(* IEC 61131-3 sources: plc-hackathon-2026/work/dump/MyController/Plc Logic/Application/Init (part 4) *)

(* ---- Init_Prof_PriceDA.st ---- *)
FUNCTION_BLOCK Init_Prof_PriceDA
VAR_INPUT
END_VAR
VAR_OUTPUT
END_VAR
VAR
END_VAR

// ---IMPL---
// Inicijalizacija GVL "Prof_PriceDA"
   Prof_PriceDA.Data[0] := 0.1353348;
   Prof_PriceDA.Data[1] := 0.1353348;
   Prof_PriceDA.Data[2] := 0.1353348;
   Prof_PriceDA.Data[3] := 0.1353348;
   Prof_PriceDA.Data[4] := 0.143694;
   Prof_PriceDA.Data[5] := 0.143694;
   Prof_PriceDA.Data[6] := 0.143694;
   Prof_PriceDA.Data[7] := 0.143694;
   Prof_PriceDA.Data[8] := 0.1349352;
   Prof_PriceDA.Data[9] := 0.1349352;
   Prof_PriceDA.Data[10] := 0.1349352;
   Prof_PriceDA.Data[11] := 0.1349352;
   Prof_PriceDA.Data[12] := 0.1010124;
   Prof_PriceDA.Data[13] := 0.1010124;
   Prof_PriceDA.Data[14] := 0.1010124;
   Prof_PriceDA.Data[15] := 0.1010124;
   Prof_PriceDA.Data[16] := 0.0687852;
   Prof_PriceDA.Data[17] := 0.0687852;
   Prof_PriceDA.Data[18] := 0.0687852;
   Prof_PriceDA.Data[19] := 0.0687852;
   Prof_PriceDA.Data[20] := 0.1011852;
   Prof_PriceDA.Data[21] := 0.1011852;
   Prof_PriceDA.Data[22] := 0.1011852;
   Prof_PriceDA.Data[23] := 0.1011852;
   Prof_PriceDA.Data[24] := 0.0974808;
   Prof_PriceDA.Data[25] := 0.0974808;
   Prof_PriceDA.Data[26] := 0.0974808;
   Prof_PriceDA.Data[27] := 0.0974808;
   Prof_PriceDA.Data[28] := 0.0902556;
   Prof_PriceDA.Data[29] := 0.0902556;
   Prof_PriceDA.Data[30] := 0.0902556;
   Prof_PriceDA.Data[31] := 0.0902556;
   Prof_PriceDA.Data[32] := 0.0399492;
   Prof_PriceDA.Data[33] := 0.0399492;
   Prof_PriceDA.Data[34] := 0.0399492;
   Prof_PriceDA.Data[35] := 0.0399492;
   Prof_PriceDA.Data[36] := 0.0485892;
   Prof_PriceDA.Data[37] := 0.0485892;
   Prof_PriceDA.Data[38] := 0.0485892;
   Prof_PriceDA.Data[39] := 0.0485892;
   Prof_PriceDA.Data[40] := 0.04158;
   Prof_PriceDA.Data[41] := 0.04158;
   Prof_PriceDA.Data[42] := 0.04158;
   Prof_PriceDA.Data[43] := 0.04158;
   Prof_PriceDA.Data[44] := 0.0430056;
   Prof_PriceDA.Data[45] := 0.0430056;
   Prof_PriceDA.Data[46] := 0.0430056;
   Prof_PriceDA.Data[47] := 0.0430056;
   Prof_PriceDA.Data[48] := 0.04347;
   Prof_PriceDA.Data[49] := 0.04347;
   Prof_PriceDA.Data[50] := 0.04347;
   Prof_PriceDA.Data[51] := 0.04347;
   Prof_PriceDA.Data[52] := 0.059886;
   Prof_PriceDA.Data[53] := 0.059886;
   Prof_PriceDA.Data[54] := 0.059886;
   Prof_PriceDA.Data[55] := 0.059886;
   Prof_PriceDA.Data[56] := 0.0664632;
   Prof_PriceDA.Data[57] := 0.0664632;
   Prof_PriceDA.Data[58] := 0.0664632;
   Prof_PriceDA.Data[59] := 0.0664632;
   Prof_PriceDA.Data[60] := 0.0900288;
   Prof_PriceDA.Data[61] := 0.0900288;
   Prof_PriceDA.Data[62] := 0.0900288;
   Prof_PriceDA.Data[63] := 0.0900288;
   Prof_PriceDA.Data[64] := 0.1161648;
   Prof_PriceDA.Data[65] := 0.1161648;
   Prof_PriceDA.Data[66] := 0.1161648;
   Prof_PriceDA.Data[67] := 0.1161648;
   Prof_PriceDA.Data[68] := 0.1328832;
   Prof_PriceDA.Data[69] := 0.1328832;
   Prof_PriceDA.Data[70] := 0.1328832;
   Prof_PriceDA.Data[71] := 0.1328832;
   Prof_PriceDA.Data[72] := 0.1382724;
   Prof_PriceDA.Data[73] := 0.1382724;
   Prof_PriceDA.Data[74] := 0.1382724;
   Prof_PriceDA.Data[75] := 0.1382724;
   Prof_PriceDA.Data[76] := 0.1446984;
   Prof_PriceDA.Data[77] := 0.1446984;
   Prof_PriceDA.Data[78] := 0.1446984;
   Prof_PriceDA.Data[79] := 0.1446984;
   Prof_PriceDA.Data[80] := 0.1406268;
   Prof_PriceDA.Data[81] := 0.1406268;
   Prof_PriceDA.Data[82] := 0.1406268;
   Prof_PriceDA.Data[83] := 0.1406268;
   Prof_PriceDA.Data[84] := 0.1307124;
   Prof_PriceDA.Data[85] := 0.1307124;
   Prof_PriceDA.Data[86] := 0.1307124;
   Prof_PriceDA.Data[87] := 0.1307124;
   Prof_PriceDA.Data[88] := 0.1310364;
   Prof_PriceDA.Data[89] := 0.1310364;
   Prof_PriceDA.Data[90] := 0.1310364;
   Prof_PriceDA.Data[91] := 0.1310364;
   Prof_PriceDA.Data[92] := 0.0904176;
   Prof_PriceDA.Data[93] := 0.0904176;
   Prof_PriceDA.Data[94] := 0.0904176;
   Prof_PriceDA.Data[95] := 0.0904176;
   Prof_PriceDA.Data[96] := 0.0689904;
   Prof_PriceDA.Data[97] := 0.0689904;
   Prof_PriceDA.Data[98] := 0.0689904;
   Prof_PriceDA.Data[99] := 0.0689904;
   Prof_PriceDA.Data[100] := 0.0865296;
   Prof_PriceDA.Data[101] := 0.0865296;
   Prof_PriceDA.Data[102] := 0.0865296;
   Prof_PriceDA.Data[103] := 0.0865296;
   Prof_PriceDA.Data[104] := 0.0846936;
   Prof_PriceDA.Data[105] := 0.0846936;
   Prof_PriceDA.Data[106] := 0.0846936;
   Prof_PriceDA.Data[107] := 0.0846936;
   Prof_PriceDA.Data[108] := 0.053136;
   Prof_PriceDA.Data[109] := 0.053136;
   Prof_PriceDA.Data[110] := 0.053136;
   Prof_PriceDA.Data[111] := 0.053136;
   Prof_PriceDA.Data[112] := 0.0614844;
   Prof_PriceDA.Data[113] := 0.0614844;
   Prof_PriceDA.Data[114] := 0.0614844;
   Prof_PriceDA.Data[115] := 0.0614844;
   Prof_PriceDA.Data[116] := 0.0834732;
   Prof_PriceDA.Data[117] := 0.0834732;
   Prof_PriceDA.Data[118] := 0.0834732;
   Prof_PriceDA.Data[119] := 0.0834732;
   Prof_PriceDA.Data[120] := 0.1200204;
   Prof_PriceDA.Data[121] := 0.1200204;
   Prof_PriceDA.Data[122] := 0.1200204;
   Prof_PriceDA.Data[123] := 0.1200204;
   Prof_PriceDA.Data[124] := 0.1431324;
   Prof_PriceDA.Data[125] := 0.1431324;
   Prof_PriceDA.Data[126] := 0.1431324;
   Prof_PriceDA.Data[127] := 0.1431324;
   Prof_PriceDA.Data[128] := 0.1405836;
   Prof_PriceDA.Data[129] := 0.1405836;
   Prof_PriceDA.Data[130] := 0.1405836;
   Prof_PriceDA.Data[131] := 0.1405836;
   Prof_PriceDA.Data[132] := 0.1433268;
   Prof_PriceDA.Data[133] := 0.1433268;
   Prof_PriceDA.Data[134] := 0.1433268;
   Prof_PriceDA.Data[135] := 0.1433268;
   Prof_PriceDA.Data[136] := 0.1391148;
   Prof_PriceDA.Data[137] := 0.1391148;
   Prof_PriceDA.Data[138] := 0.1391148;
   Prof_PriceDA.Data[139] := 0.1391148;
   Prof_PriceDA.Data[140] := 0.1337364;
   Prof_PriceDA.Data[141] := 0.1337364;
   Prof_PriceDA.Data[142] := 0.1337364;
   Prof_PriceDA.Data[143] := 0.1337364;
   Prof_PriceDA.Data[144] := 0.1330668;
   Prof_PriceDA.Data[145] := 0.1330668;
   Prof_PriceDA.Data[146] := 0.1330668;
   Prof_PriceDA.Data[147] := 0.1330668;
   Prof_PriceDA.Data[148] := 0.126144;
   Prof_PriceDA.Data[149] := 0.126144;
   Prof_PriceDA.Data[150] := 0.126144;
   Prof_PriceDA.Data[151] := 0.126144;
   Prof_PriceDA.Data[152] := 0.135;
   Prof_PriceDA.Data[153] := 0.135;
   Prof_PriceDA.Data[154] := 0.135;
   Prof_PriceDA.Data[155] := 0.135;
   Prof_PriceDA.Data[156] := 0.1405188;
   Prof_PriceDA.Data[157] := 0.1405188;
   Prof_PriceDA.Data[158] := 0.1405188;
   Prof_PriceDA.Data[159] := 0.1405188;
   Prof_PriceDA.Data[160] := 0.1650456;
   Prof_PriceDA.Data[161] := 0.1650456;
   Prof_PriceDA.Data[162] := 0.1650456;
   Prof_PriceDA.Data[163] := 0.1650456;
   Prof_PriceDA.Data[164] := 0.1762452;
   Prof_PriceDA.Data[165] := 0.1762452;
   Prof_PriceDA.Data[166] := 0.1762452;
   Prof_PriceDA.Data[167] := 0.1762452;
   Prof_PriceDA.Data[168] := 0.1695492;
   Prof_PriceDA.Data[169] := 0.1695492;
   Prof_PriceDA.Data[170] := 0.1695492;
   Prof_PriceDA.Data[171] := 0.1695492;
   Prof_PriceDA.Data[172] := 0.1646028;
   Prof_PriceDA.Data[173] := 0.1646028;
   Prof_PriceDA.Data[174] := 0.1646028;
   Prof_PriceDA.Data[175] := 0.1646028;
   Prof_PriceDA.Data[176] := 0.1414152;
   Prof_PriceDA.Data[177] := 0.1414152;
   Prof_PriceDA.Data[178] := 0.1414152;
   Prof_PriceDA.Data[179] := 0.1414152;
   Prof_PriceDA.Data[180] := 0.134622;
   Prof_PriceDA.Data[181] := 0.134622;
   Prof_PriceDA.Data[182] := 0.134622;
   Prof_PriceDA.Data[183] := 0.134622;
   Prof_PriceDA.Data[184] := 0.1270188;
   Prof_PriceDA.Data[185] := 0.1270188;
   Prof_PriceDA.Data[186] := 0.1270188;
   Prof_PriceDA.Data[187] := 0.1270188;
   Prof_PriceDA.Data[188] := 0.1095228;
   Prof_PriceDA.Data[189] := 0.1095228;
   Prof_PriceDA.Data[190] := 0.1095228;
   Prof_PriceDA.Data[191] := 0.1095228;
   Prof_PriceDA.Data[192] := 0.111996;
   Prof_PriceDA.Data[193] := 0.111996;
   Prof_PriceDA.Data[194] := 0.111996;
   Prof_PriceDA.Data[195] := 0.111996;
   Prof_PriceDA.Data[196] := 0.1023732;
   Prof_PriceDA.Data[197] := 0.1023732;
   Prof_PriceDA.Data[198] := 0.1023732;
   Prof_PriceDA.Data[199] := 0.1023732;
   Prof_PriceDA.Data[200] := 0.0968436;
   Prof_PriceDA.Data[201] := 0.0968436;
   Prof_PriceDA.Data[202] := 0.0968436;
   Prof_PriceDA.Data[203] := 0.0968436;
   Prof_PriceDA.Data[204] := 0.0945216;
   Prof_PriceDA.Data[205] := 0.0945216;
   Prof_PriceDA.Data[206] := 0.0945216;
   Prof_PriceDA.Data[207] := 0.0945216;
   Prof_PriceDA.Data[208] := 0.0923832;
   Prof_PriceDA.Data[209] := 0.0923832;
   Prof_PriceDA.Data[210] := 0.0923832;
   Prof_PriceDA.Data[211] := 0.0923832;
   Prof_PriceDA.Data[212] := 0.0993816;
   Prof_PriceDA.Data[213] := 0.0993816;
   Prof_PriceDA.Data[214] := 0.0993816;
   Prof_PriceDA.Data[215] := 0.0993816;
   Prof_PriceDA.Data[216] := 0.1185516;
   Prof_PriceDA.Data[217] := 0.1185516;
   Prof_PriceDA.Data[218] := 0.1185516;
   Prof_PriceDA.Data[219] := 0.1185516;
   Prof_PriceDA.Data[220] := 0.1469556;
   Prof_PriceDA.Data[221] := 0.1469556;
   Prof_PriceDA.Data[222] := 0.1469556;
   Prof_PriceDA.Data[223] := 0.1469556;
   Prof_PriceDA.Data[224] := 0.1492452;
   Prof_PriceDA.Data[225] := 0.1492452;
   Prof_PriceDA.Data[226] := 0.1492452;
   Prof_PriceDA.Data[227] := 0.1492452;
   Prof_PriceDA.Data[228] := 0.1461564;
   Prof_PriceDA.Data[229] := 0.1461564;
   Prof_PriceDA.Data[230] := 0.1461564;
   Prof_PriceDA.Data[231] := 0.1461564;
   Prof_PriceDA.Data[232] := 0.1350216;
   Prof_PriceDA.Data[233] := 0.1350216;
   Prof_PriceDA.Data[234] := 0.1350216;
   Prof_PriceDA.Data[235] := 0.1350216;
   Prof_PriceDA.Data[236] := 0.1219968;
   Prof_PriceDA.Data[237] := 0.1219968;
   Prof_PriceDA.Data[238] := 0.1219968;
   Prof_PriceDA.Data[239] := 0.1219968;
   Prof_PriceDA.Data[240] := 0.1201716;
   Prof_PriceDA.Data[241] := 0.1201716;
   Prof_PriceDA.Data[242] := 0.1201716;
   Prof_PriceDA.Data[243] := 0.1201716;
   Prof_PriceDA.Data[244] := 0.118206;
   Prof_PriceDA.Data[245] := 0.118206;
   Prof_PriceDA.Data[246] := 0.118206;
   Prof_PriceDA.Data[247] := 0.118206;
   Prof_PriceDA.Data[248] := 0.124956;
   Prof_PriceDA.Data[249] := 0.124956;
   Prof_PriceDA.Data[250] := 0.124956;
   Prof_PriceDA.Data[251] := 0.124956;
   Prof_PriceDA.Data[252] := 0.1402596;
   Prof_PriceDA.Data[253] := 0.1402596;
   Prof_PriceDA.Data[254] := 0.1402596;
   Prof_PriceDA.Data[255] := 0.1402596;
   Prof_PriceDA.Data[256] := 0.1587276;
   Prof_PriceDA.Data[257] := 0.1587276;
   Prof_PriceDA.Data[258] := 0.1587276;
   Prof_PriceDA.Data[259] := 0.1587276;
   Prof_PriceDA.Data[260] := 0.1571508;
   Prof_PriceDA.Data[261] := 0.1571508;
   Prof_PriceDA.Data[262] := 0.1571508;
   Prof_PriceDA.Data[263] := 0.1571508;
   Prof_PriceDA.Data[264] := 0.1572696;
   Prof_PriceDA.Data[265] := 0.1572696;
   Prof_PriceDA.Data[266] := 0.1572696;
   Prof_PriceDA.Data[267] := 0.1572696;
   Prof_PriceDA.Data[268] := 0.1564488;
   Prof_PriceDA.Data[269] := 0.1564488;
   Prof_PriceDA.Data[270] := 0.1564488;
   Prof_PriceDA.Data[271] := 0.1564488;
   Prof_PriceDA.Data[272] := 0.1478196;
   Prof_PriceDA.Data[273] := 0.1478196;
   Prof_PriceDA.Data[274] := 0.1478196;
   Prof_PriceDA.Data[275] := 0.1478196;
   Prof_PriceDA.Data[276] := 0.1314684;
   Prof_PriceDA.Data[277] := 0.1314684;
   Prof_PriceDA.Data[278] := 0.1314684;
   Prof_PriceDA.Data[279] := 0.1314684;
   Prof_PriceDA.Data[280] := 0.1361988;
   Prof_PriceDA.Data[281] := 0.1361988;
   Prof_PriceDA.Data[282] := 0.1361988;
   Prof_PriceDA.Data[283] := 0.1361988;
   Prof_PriceDA.Data[284] := 0.1318572;
   Prof_PriceDA.Data[285] := 0.1318572;
   Prof_PriceDA.Data[286] := 0.1318572;
   Prof_PriceDA.Data[287] := 0.1318572;
   Prof_PriceDA.Data[288] := 0.1189296;
   Prof_PriceDA.Data[289] := 0.1189296;
   Prof_PriceDA.Data[290] := 0.1189296;
   Prof_PriceDA.Data[291] := 0.1189296;
   Prof_PriceDA.Data[292] := 0.1130112;
   Prof_PriceDA.Data[293] := 0.1130112;
   Prof_PriceDA.Data[294] := 0.1130112;
   Prof_PriceDA.Data[295] := 0.1130112;
   Prof_PriceDA.Data[296] := 0.1087344;
   Prof_PriceDA.Data[297] := 0.1087344;
   Prof_PriceDA.Data[298] := 0.1087344;
   Prof_PriceDA.Data[299] := 0.1087344;
   Prof_PriceDA.Data[300] := 0.1065204;
   Prof_PriceDA.Data[301] := 0.1065204;
   Prof_PriceDA.Data[302] := 0.1065204;
   Prof_PriceDA.Data[303] := 0.1065204;
   Prof_PriceDA.Data[304] := 0.1077732;
   Prof_PriceDA.Data[305] := 0.1077732;
   Prof_PriceDA.Data[306] := 0.1077732;
   Prof_PriceDA.Data[307] := 0.1077732;
   Prof_PriceDA.Data[308] := 0.113454;
   Prof_PriceDA.Data[309] := 0.113454;
   Prof_PriceDA.Data[310] := 0.113454;
   Prof_PriceDA.Data[311] := 0.113454;
   Prof_PriceDA.Data[312] := 0.12096;
   Prof_PriceDA.Data[313] := 0.12096;
   Prof_PriceDA.Data[314] := 0.12096;
   Prof_PriceDA.Data[315] := 0.12096;
   Prof_PriceDA.Data[316] := 0.1352808;
   Prof_PriceDA.Data[317] := 0.1352808;
   Prof_PriceDA.Data[318] := 0.1352808;
   Prof_PriceDA.Data[319] := 0.1352808;
   Prof_PriceDA.Data[320] := 0.1386612;
   Prof_PriceDA.Data[321] := 0.1386612;
   Prof_PriceDA.Data[322] := 0.1386612;
   Prof_PriceDA.Data[323] := 0.1386612;
   Prof_PriceDA.Data[324] := 0.14121;
   Prof_PriceDA.Data[325] := 0.14121;
   Prof_PriceDA.Data[326] := 0.14121;
   Prof_PriceDA.Data[327] := 0.14121;
   Prof_PriceDA.Data[328] := 0.1407672;
   Prof_PriceDA.Data[329] := 0.1407672;
   Prof_PriceDA.Data[330] := 0.1407672;
   Prof_PriceDA.Data[331] := 0.1407672;
   Prof_PriceDA.Data[332] := 0.1385532;
   Prof_PriceDA.Data[333] := 0.1385532;
   Prof_PriceDA.Data[334] := 0.1385532;
   Prof_PriceDA.Data[335] := 0.1385532;
   Prof_PriceDA.Data[336] := 0.1404324;
   Prof_PriceDA.Data[337] := 0.1404324;
   Prof_PriceDA.Data[338] := 0.1404324;
   Prof_PriceDA.Data[339] := 0.1404324;
   Prof_PriceDA.Data[340] := 0.140238;
   Prof_PriceDA.Data[341] := 0.140238;
   Prof_PriceDA.Data[342] := 0.140238;
   Prof_PriceDA.Data[343] := 0.140238;
   Prof_PriceDA.Data[344] := 0.147312;
   Prof_PriceDA.Data[345] := 0.147312;
   Prof_PriceDA.Data[346] := 0.147312;
   Prof_PriceDA.Data[347] := 0.147312;
   Prof_PriceDA.Data[348] := 0.15309;
   Prof_PriceDA.Data[349] := 0.15309;
   Prof_PriceDA.Data[350] := 0.15309;
   Prof_PriceDA.Data[351] := 0.15309;
   Prof_PriceDA.Data[352] := 0.1819368;
   Prof_PriceDA.Data[353] := 0.1819368;
   Prof_PriceDA.Data[354] := 0.1819368;
   Prof_PriceDA.Data[355] := 0.1819368;
   Prof_PriceDA.Data[356] := 0.1857924;
   Prof_PriceDA.Data[357] := 0.1857924;
   Prof_PriceDA.Data[358] := 0.1857924;
   Prof_PriceDA.Data[359] := 0.1857924;
   Prof_PriceDA.Data[360] := 0.1848096;
   Prof_PriceDA.Data[361] := 0.1848096;
   Prof_PriceDA.Data[362] := 0.1848096;
   Prof_PriceDA.Data[363] := 0.1848096;
   Prof_PriceDA.Data[364] := 0.1831572;
   Prof_PriceDA.Data[365] := 0.1831572;
   Prof_PriceDA.Data[366] := 0.1831572;
   Prof_PriceDA.Data[367] := 0.1831572;
   Prof_PriceDA.Data[368] := 0.1590624;
   Prof_PriceDA.Data[369] := 0.1590624;
   Prof_PriceDA.Data[370] := 0.1590624;
   Prof_PriceDA.Data[371] := 0.1590624;
   Prof_PriceDA.Data[372] := 0.151524;
   Prof_PriceDA.Data[373] := 0.151524;
   Prof_PriceDA.Data[374] := 0.151524;
   Prof_PriceDA.Data[375] := 0.151524;
   Prof_PriceDA.Data[376] := 0.1455192;
   Prof_PriceDA.Data[377] := 0.1455192;
   Prof_PriceDA.Data[378] := 0.1455192;
   Prof_PriceDA.Data[379] := 0.1455192;
   Prof_PriceDA.Data[380] := 0.1259604;
   Prof_PriceDA.Data[381] := 0.1259604;
   Prof_PriceDA.Data[382] := 0.1259604;
   Prof_PriceDA.Data[383] := 0.1259604;
   Prof_PriceDA.Data[384] := 0.1211004;
   Prof_PriceDA.Data[385] := 0.1211004;
   Prof_PriceDA.Data[386] := 0.1211004;
   Prof_PriceDA.Data[387] := 0.1211004;
   Prof_PriceDA.Data[388] := 0.107838;
   Prof_PriceDA.Data[389] := 0.107838;
   Prof_PriceDA.Data[390] := 0.107838;
   Prof_PriceDA.Data[391] := 0.107838;
   Prof_PriceDA.Data[392] := 0.1033668;
   Prof_PriceDA.Data[393] := 0.1033668;
   Prof_PriceDA.Data[394] := 0.1033668;
   Prof_PriceDA.Data[395] := 0.1033668;
   Prof_PriceDA.Data[396] := 0.1013364;
   Prof_PriceDA.Data[397] := 0.1013364;
   Prof_PriceDA.Data[398] := 0.1013364;
   Prof_PriceDA.Data[399] := 0.1013364;
   Prof_PriceDA.Data[400] := 0.1006992;
   Prof_PriceDA.Data[401] := 0.1006992;
   Prof_PriceDA.Data[402] := 0.1006992;
   Prof_PriceDA.Data[403] := 0.1006992;
   Prof_PriceDA.Data[404] := 0.0971892;
   Prof_PriceDA.Data[405] := 0.0971892;
   Prof_PriceDA.Data[406] := 0.0971892;
   Prof_PriceDA.Data[407] := 0.0971892;
   Prof_PriceDA.Data[408] := 0.0989064;
   Prof_PriceDA.Data[409] := 0.0989064;
   Prof_PriceDA.Data[410] := 0.0989064;
   Prof_PriceDA.Data[411] := 0.0989064;
   Prof_PriceDA.Data[412] := 0.1068012;
   Prof_PriceDA.Data[413] := 0.1068012;
   Prof_PriceDA.Data[414] := 0.1068012;
   Prof_PriceDA.Data[415] := 0.1068012;
   Prof_PriceDA.Data[416] := 0.105408;
   Prof_PriceDA.Data[417] := 0.105408;
   Prof_PriceDA.Data[418] := 0.105408;
   Prof_PriceDA.Data[419] := 0.105408;
   Prof_PriceDA.Data[420] := 0.1070172;
   Prof_PriceDA.Data[421] := 0.1070172;
   Prof_PriceDA.Data[422] := 0.1070172;
   Prof_PriceDA.Data[423] := 0.1070172;
   Prof_PriceDA.Data[424] := 0.103194;
   Prof_PriceDA.Data[425] := 0.103194;
   Prof_PriceDA.Data[426] := 0.103194;
   Prof_PriceDA.Data[427] := 0.103194;
   Prof_PriceDA.Data[428] := 0.1084104;
   Prof_PriceDA.Data[429] := 0.1084104;
   Prof_PriceDA.Data[430] := 0.1084104;
   Prof_PriceDA.Data[431] := 0.1084104;
   Prof_PriceDA.Data[432] := 0.1057752;
   Prof_PriceDA.Data[433] := 0.1057752;
   Prof_PriceDA.Data[434] := 0.1057752;
   Prof_PriceDA.Data[435] := 0.1057752;
   Prof_PriceDA.Data[436] := 0.1129248;
   Prof_PriceDA.Data[437] := 0.1129248;
   Prof_PriceDA.Data[438] := 0.1129248;
   Prof_PriceDA.Data[439] := 0.1129248;
   Prof_PriceDA.Data[440] := 0.122094;
   Prof_PriceDA.Data[441] := 0.122094;
   Prof_PriceDA.Data[442] := 0.122094;
   Prof_PriceDA.Data[443] := 0.122094;
   Prof_PriceDA.Data[444] := 0.1337364;
   Prof_PriceDA.Data[445] := 0.1337364;
   Prof_PriceDA.Data[446] := 0.1337364;
   Prof_PriceDA.Data[447] := 0.1337364;
   Prof_PriceDA.Data[448] := 0.1717308;
   Prof_PriceDA.Data[449] := 0.1717308;
   Prof_PriceDA.Data[450] := 0.1717308;
   Prof_PriceDA.Data[451] := 0.1717308;
   Prof_PriceDA.Data[452] := 0.165024;
   Prof_PriceDA.Data[453] := 0.165024;
   Prof_PriceDA.Data[454] := 0.165024;
   Prof_PriceDA.Data[455] := 0.165024;
   Prof_PriceDA.Data[456] := 0.1562328;
   Prof_PriceDA.Data[457] := 0.1562328;
   Prof_PriceDA.Data[458] := 0.1562328;
   Prof_PriceDA.Data[459] := 0.1562328;
   Prof_PriceDA.Data[460] := 0.1627236;
   Prof_PriceDA.Data[461] := 0.1627236;
   Prof_PriceDA.Data[462] := 0.1627236;
   Prof_PriceDA.Data[463] := 0.1627236;
   Prof_PriceDA.Data[464] := 0.1535328;
   Prof_PriceDA.Data[465] := 0.1535328;
   Prof_PriceDA.Data[466] := 0.1535328;
   Prof_PriceDA.Data[467] := 0.1535328;
   Prof_PriceDA.Data[468] := 0.1449144;
   Prof_PriceDA.Data[469] := 0.1449144;
   Prof_PriceDA.Data[470] := 0.1449144;
   Prof_PriceDA.Data[471] := 0.1449144;
   Prof_PriceDA.Data[472] := 0.1105056;
   Prof_PriceDA.Data[473] := 0.1105056;
   Prof_PriceDA.Data[474] := 0.1105056;
   Prof_PriceDA.Data[475] := 0.1105056;
   Prof_PriceDA.Data[476] := 0.0771984;
   Prof_PriceDA.Data[477] := 0.0771984;
   Prof_PriceDA.Data[478] := 0.0771984;
   Prof_PriceDA.Data[479] := 0.0771984;
   Prof_PriceDA.Data[480] := 0.1130004;
   Prof_PriceDA.Data[481] := 0.1130004;
   Prof_PriceDA.Data[482] := 0.1130004;
   Prof_PriceDA.Data[483] := 0.1130004;
   Prof_PriceDA.Data[484] := 0.0960336;
   Prof_PriceDA.Data[485] := 0.0960336;
   Prof_PriceDA.Data[486] := 0.0960336;
   Prof_PriceDA.Data[487] := 0.0960336;
   Prof_PriceDA.Data[488] := 0.0743256;
   Prof_PriceDA.Data[489] := 0.0743256;
   Prof_PriceDA.Data[490] := 0.0743256;
   Prof_PriceDA.Data[491] := 0.0743256;
   Prof_PriceDA.Data[492] := 0.0708804;
   Prof_PriceDA.Data[493] := 0.0708804;
   Prof_PriceDA.Data[494] := 0.0708804;
   Prof_PriceDA.Data[495] := 0.0708804;
   Prof_PriceDA.Data[496] := 0.070794;
   Prof_PriceDA.Data[497] := 0.070794;
   Prof_PriceDA.Data[498] := 0.070794;
   Prof_PriceDA.Data[499] := 0.070794;
   Prof_PriceDA.Data[500] := 0.0962172;
   Prof_PriceDA.Data[501] := 0.0962172;
   Prof_PriceDA.Data[502] := 0.0962172;
   Prof_PriceDA.Data[503] := 0.0962172;
   Prof_PriceDA.Data[504] := 0.1229364;
   Prof_PriceDA.Data[505] := 0.1229364;
   Prof_PriceDA.Data[506] := 0.1229364;
   Prof_PriceDA.Data[507] := 0.1229364;
   Prof_PriceDA.Data[508] := 0.1331748;
   Prof_PriceDA.Data[509] := 0.1331748;
   Prof_PriceDA.Data[510] := 0.1331748;
   Prof_PriceDA.Data[511] := 0.1331748;
   Prof_PriceDA.Data[512] := 0.1334664;
   Prof_PriceDA.Data[513] := 0.1334664;
   Prof_PriceDA.Data[514] := 0.1334664;
   Prof_PriceDA.Data[515] := 0.1334664;
   Prof_PriceDA.Data[516] := 0.1152576;
   Prof_PriceDA.Data[517] := 0.1152576;
   Prof_PriceDA.Data[518] := 0.1152576;
   Prof_PriceDA.Data[519] := 0.1152576;
   Prof_PriceDA.Data[520] := 0.097956;
   Prof_PriceDA.Data[521] := 0.097956;
   Prof_PriceDA.Data[522] := 0.097956;
   Prof_PriceDA.Data[523] := 0.097956;
   Prof_PriceDA.Data[524] := 0.0780624;
   Prof_PriceDA.Data[525] := 0.0780624;
   Prof_PriceDA.Data[526] := 0.0780624;
   Prof_PriceDA.Data[527] := 0.0780624;
   Prof_PriceDA.Data[528] := 0.0841212;
   Prof_PriceDA.Data[529] := 0.0841212;
   Prof_PriceDA.Data[530] := 0.0841212;
   Prof_PriceDA.Data[531] := 0.0841212;
   Prof_PriceDA.Data[532] := 0.10476;
   Prof_PriceDA.Data[533] := 0.10476;
   Prof_PriceDA.Data[534] := 0.10476;
   Prof_PriceDA.Data[535] := 0.10476;
   Prof_PriceDA.Data[536] := 0.1249668;
   Prof_PriceDA.Data[537] := 0.1249668;
   Prof_PriceDA.Data[538] := 0.1249668;
   Prof_PriceDA.Data[539] := 0.1249668;
   Prof_PriceDA.Data[540] := 0.1229904;
   Prof_PriceDA.Data[541] := 0.1229904;
   Prof_PriceDA.Data[542] := 0.1229904;
   Prof_PriceDA.Data[543] := 0.1229904;
   Prof_PriceDA.Data[544] := 0.1472904;
   Prof_PriceDA.Data[545] := 0.1472904;
   Prof_PriceDA.Data[546] := 0.1472904;
   Prof_PriceDA.Data[547] := 0.1472904;
   Prof_PriceDA.Data[548] := 0.1600344;
   Prof_PriceDA.Data[549] := 0.1600344;
   Prof_PriceDA.Data[550] := 0.1600344;
   Prof_PriceDA.Data[551] := 0.1600344;
   Prof_PriceDA.Data[552] := 0.1528524;
   Prof_PriceDA.Data[553] := 0.1528524;
   Prof_PriceDA.Data[554] := 0.1528524;
   Prof_PriceDA.Data[555] := 0.1528524;
   Prof_PriceDA.Data[556] := 0.1521828;
   Prof_PriceDA.Data[557] := 0.1521828;
   Prof_PriceDA.Data[558] := 0.1521828;
   Prof_PriceDA.Data[559] := 0.1521828;
   Prof_PriceDA.Data[560] := 0.1456272;
   Prof_PriceDA.Data[561] := 0.1456272;
   Prof_PriceDA.Data[562] := 0.1456272;
   Prof_PriceDA.Data[563] := 0.1456272;
   Prof_PriceDA.Data[564] := 0.122364;
   Prof_PriceDA.Data[565] := 0.122364;
   Prof_PriceDA.Data[566] := 0.122364;
   Prof_PriceDA.Data[567] := 0.122364;
   Prof_PriceDA.Data[568] := 0.1168128;
   Prof_PriceDA.Data[569] := 0.1168128;
   Prof_PriceDA.Data[570] := 0.1168128;
   Prof_PriceDA.Data[571] := 0.1168128;
   Prof_PriceDA.Data[572] := 0.0853416;
   Prof_PriceDA.Data[573] := 0.0853416;
   Prof_PriceDA.Data[574] := 0.0853416;
   Prof_PriceDA.Data[575] := 0.0853416;
   Prof_PriceDA.Data[576] := 0.0343116;
   Prof_PriceDA.Data[577] := 0.0343116;
   Prof_PriceDA.Data[578] := 0.0343116;
   Prof_PriceDA.Data[579] := 0.0343116;
   Prof_PriceDA.Data[580] := 0.056538;
   Prof_PriceDA.Data[581] := 0.056538;
   Prof_PriceDA.Data[582] := 0.056538;
   Prof_PriceDA.Data[583] := 0.056538;
   Prof_PriceDA.Data[584] := 0.0510192;
   Prof_PriceDA.Data[585] := 0.0510192;
   Prof_PriceDA.Data[586] := 0.0510192;
   Prof_PriceDA.Data[587] := 0.0510192;
   Prof_PriceDA.Data[588] := 0.0135;
   Prof_PriceDA.Data[589] := 0.0135;
   Prof_PriceDA.Data[590] := 0.0135;
   Prof_PriceDA.Data[591] := 0.0135;
   Prof_PriceDA.Data[592] := 0.0662688;
   Prof_PriceDA.Data[593] := 0.0662688;
   Prof_PriceDA.Data[594] := 0.0662688;
   Prof_PriceDA.Data[595] := 0.0662688;
   Prof_PriceDA.Data[596] := 0.0844668;
   Prof_PriceDA.Data[597] := 0.0844668;
   Prof_PriceDA.Data[598] := 0.0844668;
   Prof_PriceDA.Data[599] := 0.0844668;
   Prof_PriceDA.Data[600] := 0.1362636;
   Prof_PriceDA.Data[601] := 0.1362636;
   Prof_PriceDA.Data[602] := 0.1362636;
   Prof_PriceDA.Data[603] := 0.1362636;
   Prof_PriceDA.Data[604] := 0.16443;
   Prof_PriceDA.Data[605] := 0.16443;
   Prof_PriceDA.Data[606] := 0.16443;
   Prof_PriceDA.Data[607] := 0.16443;
   Prof_PriceDA.Data[608] := 0.148014;
   Prof_PriceDA.Data[609] := 0.148014;
   Prof_PriceDA.Data[610] := 0.148014;
   Prof_PriceDA.Data[611] := 0.148014;
   Prof_PriceDA.Data[612] := 0.1423224;
   Prof_PriceDA.Data[613] := 0.1423224;
   Prof_PriceDA.Data[614] := 0.1423224;
   Prof_PriceDA.Data[615] := 0.1423224;
   Prof_PriceDA.Data[616] := 0.1318248;
   Prof_PriceDA.Data[617] := 0.1318248;
   Prof_PriceDA.Data[618] := 0.1318248;
   Prof_PriceDA.Data[619] := 0.1318248;
   Prof_PriceDA.Data[620] := 0.131274;
   Prof_PriceDA.Data[621] := 0.131274;
   Prof_PriceDA.Data[622] := 0.131274;
   Prof_PriceDA.Data[623] := 0.131274;
   Prof_PriceDA.Data[624] := 0.1322676;
   Prof_PriceDA.Data[625] := 0.1322676;
   Prof_PriceDA.Data[626] := 0.1322676;
   Prof_PriceDA.Data[627] := 0.1322676;
   Prof_PriceDA.Data[628] := 0.1404432;
   Prof_PriceDA.Data[629] := 0.1404432;
   Prof_PriceDA.Data[630] := 0.1404432;
   Prof_PriceDA.Data[631] := 0.1404432;
   Prof_PriceDA.Data[632] := 0.1504656;
   Prof_PriceDA.Data[633] := 0.1504656;
   Prof_PriceDA.Data[634] := 0.1504656;
   Prof_PriceDA.Data[635] := 0.1504656;
   Prof_PriceDA.Data[636] := 0.1588572;
   Prof_PriceDA.Data[637] := 0.1588572;
   Prof_PriceDA.Data[638] := 0.1588572;
   Prof_PriceDA.Data[639] := 0.1588572;
   Prof_PriceDA.Data[640] := 0.1668384;
   Prof_PriceDA.Data[641] := 0.1668384;
   Prof_PriceDA.Data[642] := 0.1668384;
   Prof_PriceDA.Data[643] := 0.1668384;
   Prof_PriceDA.Data[644] := 0.166806;
   Prof_PriceDA.Data[645] := 0.166806;
   Prof_PriceDA.Data[646] := 0.166806;
   Prof_PriceDA.Data[647] := 0.166806;
   Prof_PriceDA.Data[648] := 0.1628424;
   Prof_PriceDA.Data[649] := 0.1628424;
   Prof_PriceDA.Data[650] := 0.1628424;
   Prof_PriceDA.Data[651] := 0.1628424;
   Prof_PriceDA.Data[652] := 0.1643328;
   Prof_PriceDA.Data[653] := 0.1643328;
   Prof_PriceDA.Data[654] := 0.1643328;
   Prof_PriceDA.Data[655] := 0.1643328;
   Prof_PriceDA.Data[656] := 0.1532088;
   Prof_PriceDA.Data[657] := 0.1532088;
   Prof_PriceDA.Data[658] := 0.1532088;
   Prof_PriceDA.Data[659] := 0.1532088;
   Prof_PriceDA.Data[660] := 0.1370196;
   Prof_PriceDA.Data[661] := 0.1370196;
   Prof_PriceDA.Data[662] := 0.1370196;
   Prof_PriceDA.Data[663] := 0.1370196;
   Prof_PriceDA.Data[664] := 0.125064;
   Prof_PriceDA.Data[665] := 0.125064;
   Prof_PriceDA.Data[666] := 0.125064;
   Prof_PriceDA.Data[667] := 0.125064;
   Prof_PriceDA.Data[668] := 0.1204416;
   Prof_PriceDA.Data[669] := 0.1204416;
   Prof_PriceDA.Data[670] := 0.1204416;
   Prof_PriceDA.Data[671] := 0.1204416;
   Prof_PriceDA.Data[672] := 0.0901584;
   Prof_PriceDA.Data[673] := 0.0901584;
   Prof_PriceDA.Data[674] := 0.0901584;
   Prof_PriceDA.Data[675] := 0.0901584;
   Prof_PriceDA.Data[676] := 0.0813672;
   Prof_PriceDA.Data[677] := 0.0813672;
   Prof_PriceDA.Data[678] := 0.0813672;
   Prof_PriceDA.Data[679] := 0.0813672;
   Prof_PriceDA.Data[680] := 0.0789048;
   Prof_PriceDA.Data[681] := 0.0789048;
   Prof_PriceDA.Data[682] := 0.0789048;
   Prof_PriceDA.Data[683] := 0.0789048;
   Prof_PriceDA.Data[684] := 0.0747036;
   Prof_PriceDA.Data[685] := 0.0747036;
   Prof_PriceDA.Data[686] := 0.0747036;
   Prof_PriceDA.Data[687] := 0.0747036;
   Prof_PriceDA.Data[688] := 0.0923076;
   Prof_PriceDA.Data[689] := 0.0923076;
   Prof_PriceDA.Data[690] := 0.0923076;
   Prof_PriceDA.Data[691] := 0.0923076;
   Prof_PriceDA.Data[692] := 0.11178;
   Prof_PriceDA.Data[693] := 0.11178;
   Prof_PriceDA.Data[694] := 0.11178;
   Prof_PriceDA.Data[695] := 0.11178;
   Prof_PriceDA.Data[696] := 0.1367388;
   Prof_PriceDA.Data[697] := 0.1367388;
   Prof_PriceDA.Data[698] := 0.1367388;
   Prof_PriceDA.Data[699] := 0.1367388;
   Prof_PriceDA.Data[700] := 0.1635336;
   Prof_PriceDA.Data[701] := 0.1635336;
   Prof_PriceDA.Data[702] := 0.1635336;
   Prof_PriceDA.Data[703] := 0.1635336;
   Prof_PriceDA.Data[704] := 0.1611252;
   Prof_PriceDA.Data[705] := 0.1611252;
   Prof_PriceDA.Data[706] := 0.1611252;
   Prof_PriceDA.Data[707] := 0.1611252;
   Prof_PriceDA.Data[708] := 0.1341576;
   Prof_PriceDA.Data[709] := 0.1341576;
   Prof_PriceDA.Data[710] := 0.1341576;
   Prof_PriceDA.Data[711] := 0.1341576;
   Prof_PriceDA.Data[712] := 0.1174068;
   Prof_PriceDA.Data[713] := 0.1174068;
   Prof_PriceDA.Data[714] := 0.1174068;
   Prof_PriceDA.Data[715] := 0.1174068;
   Prof_PriceDA.Data[716] := 0.1103436;
   Prof_PriceDA.Data[717] := 0.1103436;
   Prof_PriceDA.Data[718] := 0.1103436;
   Prof_PriceDA.Data[719] := 0.1103436;
   Prof_PriceDA.Data[720] := 0.1120824;
   Prof_PriceDA.Data[721] := 0.1120824;
   Prof_PriceDA.Data[722] := 0.1120824;
   Prof_PriceDA.Data[723] := 0.1120824;
   Prof_PriceDA.Data[724] := 0.1245996;
   Prof_PriceDA.Data[725] := 0.1245996;
   Prof_PriceDA.Data[726] := 0.1245996;
   Prof_PriceDA.Data[727] := 0.1245996;
   Prof_PriceDA.Data[728] := 0.1353132;
   Prof_PriceDA.Data[729] := 0.1353132;
   Prof_PriceDA.Data[730] := 0.1353132;
   Prof_PriceDA.Data[731] := 0.1353132;
   Prof_PriceDA.Data[732] := 0.1550556;
   Prof_PriceDA.Data[733] := 0.1550556;
   Prof_PriceDA.Data[734] := 0.1550556;
   Prof_PriceDA.Data[735] := 0.1550556;
   Prof_PriceDA.Data[736] := 0.1646784;
   Prof_PriceDA.Data[737] := 0.1646784;
   Prof_PriceDA.Data[738] := 0.1646784;
   Prof_PriceDA.Data[739] := 0.1646784;
   Prof_PriceDA.Data[740] := 0.165456;
   Prof_PriceDA.Data[741] := 0.165456;
   Prof_PriceDA.Data[742] := 0.165456;
   Prof_PriceDA.Data[743] := 0.165456;
   Prof_PriceDA.Data[744] := 0.1622916;
   Prof_PriceDA.Data[745] := 0.1622916;
   Prof_PriceDA.Data[746] := 0.1622916;
   Prof_PriceDA.Data[747] := 0.1622916;
   Prof_PriceDA.Data[748] := 0.1614384;
   Prof_PriceDA.Data[749] := 0.1614384;
   Prof_PriceDA.Data[750] := 0.1614384;
   Prof_PriceDA.Data[751] := 0.1614384;
   Prof_PriceDA.Data[752] := 0.1484352;
   Prof_PriceDA.Data[753] := 0.1484352;
   Prof_PriceDA.Data[754] := 0.1484352;
   Prof_PriceDA.Data[755] := 0.1484352;
   Prof_PriceDA.Data[756] := 0.1356372;
   Prof_PriceDA.Data[757] := 0.1356372;
   Prof_PriceDA.Data[758] := 0.1356372;
   Prof_PriceDA.Data[759] := 0.1356372;
   Prof_PriceDA.Data[760] := 0.1255716;
   Prof_PriceDA.Data[761] := 0.1255716;
   Prof_PriceDA.Data[762] := 0.1255716;
   Prof_PriceDA.Data[763] := 0.1255716;
   Prof_PriceDA.Data[764] := 0.114588;
   Prof_PriceDA.Data[765] := 0.114588;
   Prof_PriceDA.Data[766] := 0.114588;
   Prof_PriceDA.Data[767] := 0.114588;
   Prof_PriceDA.Data[768] := 0.1147284;
   Prof_PriceDA.Data[769] := 0.1147284;
   Prof_PriceDA.Data[770] := 0.1147284;
   Prof_PriceDA.Data[771] := 0.1147284;
   Prof_PriceDA.Data[772] := 0.114588;
   Prof_PriceDA.Data[773] := 0.114588;
   Prof_PriceDA.Data[774] := 0.114588;
   Prof_PriceDA.Data[775] := 0.114588;
   Prof_PriceDA.Data[776] := 0.1119096;
   Prof_PriceDA.Data[777] := 0.1119096;
   Prof_PriceDA.Data[778] := 0.1119096;
   Prof_PriceDA.Data[779] := 0.1119096;
   Prof_PriceDA.Data[780] := 0.1104408;
   Prof_PriceDA.Data[781] := 0.1104408;
   Prof_PriceDA.Data[782] := 0.1104408;
   Prof_PriceDA.Data[783] := 0.1104408;
   Prof_PriceDA.Data[784] := 0.1152468;
   Prof_PriceDA.Data[785] := 0.1152468;
   Prof_PriceDA.Data[786] := 0.1152468;
   Prof_PriceDA.Data[787] := 0.1152468;
   Prof_PriceDA.Data[788] := 0.1184868;
   Prof_PriceDA.Data[789] := 0.1184868;
   Prof_PriceDA.Data[790] := 0.1184868;
   Prof_PriceDA.Data[791] := 0.1184868;
   Prof_PriceDA.Data[792] := 0.1342656;
   Prof_PriceDA.Data[793] := 0.1342656;
   Prof_PriceDA.Data[794] := 0.1342656;
   Prof_PriceDA.Data[795] := 0.1342656;
   Prof_PriceDA.Data[796] := 0.1542132;
   Prof_PriceDA.Data[797] := 0.1542132;
   Prof_PriceDA.Data[798] := 0.1542132;
   Prof_PriceDA.Data[799] := 0.1542132;
   Prof_PriceDA.Data[800] := 0.1678104;
   Prof_PriceDA.Data[801] := 0.1678104;
   Prof_PriceDA.Data[802] := 0.1678104;
   Prof_PriceDA.Data[803] := 0.1678104;
   Prof_PriceDA.Data[804] := 0.1601208;
   Prof_PriceDA.Data[805] := 0.1601208;
   Prof_PriceDA.Data[806] := 0.1601208;
   Prof_PriceDA.Data[807] := 0.1601208;
   Prof_PriceDA.Data[808] := 0.1514916;
   Prof_PriceDA.Data[809] := 0.1514916;
   Prof_PriceDA.Data[810] := 0.1514916;
   Prof_PriceDA.Data[811] := 0.1514916;
   Prof_PriceDA.Data[812] := 0.1435644;
   Prof_PriceDA.Data[813] := 0.1435644;
   Prof_PriceDA.Data[814] := 0.1435644;
   Prof_PriceDA.Data[815] := 0.1435644;
   Prof_PriceDA.Data[816] := 0.1331532;
   Prof_PriceDA.Data[817] := 0.1331532;
   Prof_PriceDA.Data[818] := 0.1331532;
   Prof_PriceDA.Data[819] := 0.1331532;
   Prof_PriceDA.Data[820] := 0.1284012;
   Prof_PriceDA.Data[821] := 0.1284012;
   Prof_PriceDA.Data[822] := 0.1284012;
   Prof_PriceDA.Data[823] := 0.1284012;
   Prof_PriceDA.Data[824] := 0.1325484;
   Prof_PriceDA.Data[825] := 0.1325484;
   Prof_PriceDA.Data[826] := 0.1325484;
   Prof_PriceDA.Data[827] := 0.1325484;
   Prof_PriceDA.Data[828] := 0.1425708;
   Prof_PriceDA.Data[829] := 0.1425708;
   Prof_PriceDA.Data[830] := 0.1425708;
   Prof_PriceDA.Data[831] := 0.1425708;
   Prof_PriceDA.Data[832] := 0.1583496;
   Prof_PriceDA.Data[833] := 0.1583496;
   Prof_PriceDA.Data[834] := 0.1583496;
   Prof_PriceDA.Data[835] := 0.1583496;
   Prof_PriceDA.Data[836] := 0.1566756;
   Prof_PriceDA.Data[837] := 0.1566756;
   Prof_PriceDA.Data[838] := 0.1566756;
   Prof_PriceDA.Data[839] := 0.1566756;
   Prof_PriceDA.Data[840] := 0.16065;
   Prof_PriceDA.Data[841] := 0.16065;
   Prof_PriceDA.Data[842] := 0.16065;
   Prof_PriceDA.Data[843] := 0.16065;
   Prof_PriceDA.Data[844] := 0.1521612;
   Prof_PriceDA.Data[845] := 0.1521612;
   Prof_PriceDA.Data[846] := 0.1521612;
   Prof_PriceDA.Data[847] := 0.1521612;
   Prof_PriceDA.Data[848] := 0.1421172;
   Prof_PriceDA.Data[849] := 0.1421172;
   Prof_PriceDA.Data[850] := 0.1421172;
   Prof_PriceDA.Data[851] := 0.1421172;
   Prof_PriceDA.Data[852] := 0.1240056;
   Prof_PriceDA.Data[853] := 0.1240056;
   Prof_PriceDA.Data[854] := 0.1240056;
   Prof_PriceDA.Data[855] := 0.1240056;
   Prof_PriceDA.Data[856] := 0.11151;
   Prof_PriceDA.Data[857] := 0.11151;
   Prof_PriceDA.Data[858] := 0.11151;
   Prof_PriceDA.Data[859] := 0.11151;
   Prof_PriceDA.Data[860] := 0.0968328;
   Prof_PriceDA.Data[861] := 0.0968328;
   Prof_PriceDA.Data[862] := 0.0968328;
   Prof_PriceDA.Data[863] := 0.0968328;
   Prof_PriceDA.Data[864] := 0.0941976;
   Prof_PriceDA.Data[865] := 0.0941976;
   Prof_PriceDA.Data[866] := 0.0941976;
   Prof_PriceDA.Data[867] := 0.0941976;
   Prof_PriceDA.Data[868] := 0.0868104;
   Prof_PriceDA.Data[869] := 0.0868104;
   Prof_PriceDA.Data[870] := 0.0868104;
   Prof_PriceDA.Data[871] := 0.0868104;
   Prof_PriceDA.Data[872] := 0.0826092;
   Prof_PriceDA.Data[873] := 0.0826092;
   Prof_PriceDA.Data[874] := 0.0826092;
   Prof_PriceDA.Data[875] := 0.0826092;
   Prof_PriceDA.Data[876] := 0.0808164;
   Prof_PriceDA.Data[877] := 0.0808164;
   Prof_PriceDA.Data[878] := 0.0808164;
   Prof_PriceDA.Data[879] := 0.0808164;
   Prof_PriceDA.Data[880] := 0.0767664;
   Prof_PriceDA.Data[881] := 0.0767664;
   Prof_PriceDA.Data[882] := 0.0767664;
   Prof_PriceDA.Data[883] := 0.0767664;
   Prof_PriceDA.Data[884] := 0.1046088;
   Prof_PriceDA.Data[885] := 0.1046088;
   Prof_PriceDA.Data[886] := 0.1046088;
   Prof_PriceDA.Data[887] := 0.1046088;
   Prof_PriceDA.Data[888] := 0.1354968;
   Prof_PriceDA.Data[889] := 0.1354968;
   Prof_PriceDA.Data[890] := 0.1354968;
   Prof_PriceDA.Data[891] := 0.1354968;
   Prof_PriceDA.Data[892] := 0.165024;
   Prof_PriceDA.Data[893] := 0.165024;
   Prof_PriceDA.Data[894] := 0.165024;
   Prof_PriceDA.Data[895] := 0.165024;
   Prof_PriceDA.Data[896] := 0.1680264;
   Prof_PriceDA.Data[897] := 0.1680264;
   Prof_PriceDA.Data[898] := 0.1680264;
   Prof_PriceDA.Data[899] := 0.1680264;
   Prof_PriceDA.Data[900] := 0.1522368;
   Prof_PriceDA.Data[901] := 0.1522368;
   Prof_PriceDA.Data[902] := 0.1522368;
   Prof_PriceDA.Data[903] := 0.1522368;
   Prof_PriceDA.Data[904] := 0.1334556;
   Prof_PriceDA.Data[905] := 0.1334556;
   Prof_PriceDA.Data[906] := 0.1334556;
   Prof_PriceDA.Data[907] := 0.1334556;
   Prof_PriceDA.Data[908] := 0.1226772;
   Prof_PriceDA.Data[909] := 0.1226772;
   Prof_PriceDA.Data[910] := 0.1226772;
   Prof_PriceDA.Data[911] := 0.1226772;
   Prof_PriceDA.Data[912] := 0.1160244;
   Prof_PriceDA.Data[913] := 0.1160244;
   Prof_PriceDA.Data[914] := 0.1160244;
   Prof_PriceDA.Data[915] := 0.1160244;
   Prof_PriceDA.Data[916] := 0.1134108;
   Prof_PriceDA.Data[917] := 0.1134108;
   Prof_PriceDA.Data[918] := 0.1134108;
   Prof_PriceDA.Data[919] := 0.1134108;
   Prof_PriceDA.Data[920] := 0.1188108;
   Prof_PriceDA.Data[921] := 0.1188108;
   Prof_PriceDA.Data[922] := 0.1188108;
   Prof_PriceDA.Data[923] := 0.1188108;
   Prof_PriceDA.Data[924] := 0.1389852;
   Prof_PriceDA.Data[925] := 0.1389852;
   Prof_PriceDA.Data[926] := 0.1389852;
   Prof_PriceDA.Data[927] := 0.1389852;
   Prof_PriceDA.Data[928] := 0.1609308;
   Prof_PriceDA.Data[929] := 0.1609308;
   Prof_PriceDA.Data[930] := 0.1609308;
   Prof_PriceDA.Data[931] := 0.1609308;
   Prof_PriceDA.Data[932] := 0.1583604;
   Prof_PriceDA.Data[933] := 0.1583604;
   Prof_PriceDA.Data[934] := 0.1583604;
   Prof_PriceDA.Data[935] := 0.1583604;
   Prof_PriceDA.Data[936] := 0.1590084;
   Prof_PriceDA.Data[937] := 0.1590084;
   Prof_PriceDA.Data[938] := 0.1590084;
   Prof_PriceDA.Data[939] := 0.1590084;
   Prof_PriceDA.Data[940] := 0.1569024;
   Prof_PriceDA.Data[941] := 0.1569024;
   Prof_PriceDA.Data[942] := 0.1569024;
   Prof_PriceDA.Data[943] := 0.1569024;
   Prof_PriceDA.Data[944] := 0.1457568;
   Prof_PriceDA.Data[945] := 0.1457568;
   Prof_PriceDA.Data[946] := 0.1457568;
   Prof_PriceDA.Data[947] := 0.1457568;
   Prof_PriceDA.Data[948] := 0.1323108;
   Prof_PriceDA.Data[949] := 0.1323108;
   Prof_PriceDA.Data[950] := 0.1323108;
   Prof_PriceDA.Data[951] := 0.1323108;
   Prof_PriceDA.Data[952] := 0.129492;
   Prof_PriceDA.Data[953] := 0.129492;
   Prof_PriceDA.Data[954] := 0.129492;
   Prof_PriceDA.Data[955] := 0.129492;
   Prof_PriceDA.Data[956] := 0.1226016;
   Prof_PriceDA.Data[957] := 0.1226016;
   Prof_PriceDA.Data[958] := 0.1226016;
   Prof_PriceDA.Data[959] := 0.1226016;
   Prof_PriceDA.Data[960] := 0.1179468;
   Prof_PriceDA.Data[961] := 0.1179468;
   Prof_PriceDA.Data[962] := 0.1179468;
   Prof_PriceDA.Data[963] := 0.1179468;
   Prof_PriceDA.Data[964] := 0.1079676;
   Prof_PriceDA.Data[965] := 0.1079676;
   Prof_PriceDA.Data[966] := 0.1079676;
   Prof_PriceDA.Data[967] := 0.1079676;
   Prof_PriceDA.Data[968] := 0.1042632;
   Prof_PriceDA.Data[969] := 0.1042632;
   Prof_PriceDA.Data[970] := 0.1042632;
   Prof_PriceDA.Data[971] := 0.1042632;
   Prof_PriceDA.Data[972] := 0.1000296;
   Prof_PriceDA.Data[973] := 0.1000296;
   Prof_PriceDA.Data[974] := 0.1000296;
   Prof_PriceDA.Data[975] := 0.1000296;
   Prof_PriceDA.Data[976] := 0.099144;
   Prof_PriceDA.Data[977] := 0.099144;
   Prof_PriceDA.Data[978] := 0.099144;
   Prof_PriceDA.Data[979] := 0.099144;
   Prof_PriceDA.Data[980] := 0.1006236;
   Prof_PriceDA.Data[981] := 0.1006236;
   Prof_PriceDA.Data[982] := 0.1006236;
   Prof_PriceDA.Data[983] := 0.1006236;
   Prof_PriceDA.Data[984] := 0.1021788;
   Prof_PriceDA.Data[985] := 0.1021788;
   Prof_PriceDA.Data[986] := 0.1021788;
   Prof_PriceDA.Data[987] := 0.1021788;
   Prof_PriceDA.Data[988] := 0.1209168;
   Prof_PriceDA.Data[989] := 0.1209168;
   Prof_PriceDA.Data[990] := 0.1209168;
   Prof_PriceDA.Data[991] := 0.1209168;
   Prof_PriceDA.Data[992] := 0.12312;
   Prof_PriceDA.Data[993] := 0.12312;
   Prof_PriceDA.Data[994] := 0.12312;
   Prof_PriceDA.Data[995] := 0.12312;
   Prof_PriceDA.Data[996] := 0.1200744;
   Prof_PriceDA.Data[997] := 0.1200744;
   Prof_PriceDA.Data[998] := 0.1200744;
   Prof_PriceDA.Data[999] := 0.1200744;
   Prof_PriceDA.Data[1000] := 0.113454;
   Prof_PriceDA.Data[1001] := 0.113454;
   Prof_PriceDA.Data[1002] := 0.113454;
   Prof_PriceDA.Data[1003] := 0.113454;
   Prof_PriceDA.Data[1004] := 0.1078488;
   Prof_PriceDA.Data[1005] := 0.1078488;
   Prof_PriceDA.Data[1006] := 0.1078488;
   Prof_PriceDA.Data[1007] := 0.1078488;
   Prof_PriceDA.Data[1008] := 0.1046088;
   Prof_PriceDA.Data[1009] := 0.1046088;
   Prof_PriceDA.Data[1010] := 0.1046088;
   Prof_PriceDA.Data[1011] := 0.1046088;
   Prof_PriceDA.Data[1012] := 0.100602;
   Prof_PriceDA.Data[1013] := 0.100602;
   Prof_PriceDA.Data[1014] := 0.100602;
   Prof_PriceDA.Data[1015] := 0.100602;
   Prof_PriceDA.Data[1016] := 0.1068768;
   Prof_PriceDA.Data[1017] := 0.1068768;
   Prof_PriceDA.Data[1018] := 0.1068768;
   Prof_PriceDA.Data[1019] := 0.1068768;
   Prof_PriceDA.Data[1020] := 0.113994;
   Prof_PriceDA.Data[1021] := 0.113994;
   Prof_PriceDA.Data[1022] := 0.113994;
   Prof_PriceDA.Data[1023] := 0.113994;
   Prof_PriceDA.Data[1024] := 0.1448928;
   Prof_PriceDA.Data[1025] := 0.1448928;
   Prof_PriceDA.Data[1026] := 0.1448928;
   Prof_PriceDA.Data[1027] := 0.1448928;
   Prof_PriceDA.Data[1028] := 0.1509732;
   Prof_PriceDA.Data[1029] := 0.1509732;
   Prof_PriceDA.Data[1030] := 0.1509732;
   Prof_PriceDA.Data[1031] := 0.1509732;
   Prof_PriceDA.Data[1032] := 0.1472256;
   Prof_PriceDA.Data[1033] := 0.1472256;
   Prof_PriceDA.Data[1034] := 0.1472256;
   Prof_PriceDA.Data[1035] := 0.1472256;
   Prof_PriceDA.Data[1036] := 0.148284;
   Prof_PriceDA.Data[1037] := 0.148284;
   Prof_PriceDA.Data[1038] := 0.148284;
   Prof_PriceDA.Data[1039] := 0.148284;
   Prof_PriceDA.Data[1040] := 0.1366848;
   Prof_PriceDA.Data[1041] := 0.1366848;
   Prof_PriceDA.Data[1042] := 0.1366848;
   Prof_PriceDA.Data[1043] := 0.1366848;
   Prof_PriceDA.Data[1044] := 0.1265328;
   Prof_PriceDA.Data[1045] := 0.1265328;
   Prof_PriceDA.Data[1046] := 0.1265328;
   Prof_PriceDA.Data[1047] := 0.1265328;
   Prof_PriceDA.Data[1048] := 0.11799;
   Prof_PriceDA.Data[1049] := 0.11799;
   Prof_PriceDA.Data[1050] := 0.11799;
   Prof_PriceDA.Data[1051] := 0.11799;
   Prof_PriceDA.Data[1052] := 0.1143612;
   Prof_PriceDA.Data[1053] := 0.1143612;
   Prof_PriceDA.Data[1054] := 0.1143612;
   Prof_PriceDA.Data[1055] := 0.1143612;
   Prof_PriceDA.Data[1056] := 0.1075896;
   Prof_PriceDA.Data[1057] := 0.1075896;
   Prof_PriceDA.Data[1058] := 0.1075896;
   Prof_PriceDA.Data[1059] := 0.1075896;
   Prof_PriceDA.Data[1060] := 0.0961416;
   Prof_PriceDA.Data[1061] := 0.0961416;
   Prof_PriceDA.Data[1062] := 0.0961416;
   Prof_PriceDA.Data[1063] := 0.0961416;
   Prof_PriceDA.Data[1064] := 0.0964548;
   Prof_PriceDA.Data[1065] := 0.0964548;
   Prof_PriceDA.Data[1066] := 0.0964548;
   Prof_PriceDA.Data[1067] := 0.0964548;
   Prof_PriceDA.Data[1068] := 0.092178;
   Prof_PriceDA.Data[1069] := 0.092178;
   Prof_PriceDA.Data[1070] := 0.092178;
   Prof_PriceDA.Data[1071] := 0.092178;
   Prof_PriceDA.Data[1072] := 0.0918;
   Prof_PriceDA.Data[1073] := 0.0918;
   Prof_PriceDA.Data[1074] := 0.0918;
   Prof_PriceDA.Data[1075] := 0.0918;
   Prof_PriceDA.Data[1076] := 0.0919188;
   Prof_PriceDA.Data[1077] := 0.0919188;
   Prof_PriceDA.Data[1078] := 0.0919188;
   Prof_PriceDA.Data[1079] := 0.0919188;
   Prof_PriceDA.Data[1080] := 0.0946836;
   Prof_PriceDA.Data[1081] := 0.0946836;
   Prof_PriceDA.Data[1082] := 0.0946836;
   Prof_PriceDA.Data[1083] := 0.0946836;
   Prof_PriceDA.Data[1084] := 0.10989;
   Prof_PriceDA.Data[1085] := 0.10989;
   Prof_PriceDA.Data[1086] := 0.10989;
   Prof_PriceDA.Data[1087] := 0.10989;
   Prof_PriceDA.Data[1088] := 0.1258092;
   Prof_PriceDA.Data[1089] := 0.1258092;
   Prof_PriceDA.Data[1090] := 0.1258092;
   Prof_PriceDA.Data[1091] := 0.1258092;
   Prof_PriceDA.Data[1092] := 0.1296756;
   Prof_PriceDA.Data[1093] := 0.1296756;
   Prof_PriceDA.Data[1094] := 0.1296756;
   Prof_PriceDA.Data[1095] := 0.1296756;
   Prof_PriceDA.Data[1096] := 0.1271916;
   Prof_PriceDA.Data[1097] := 0.1271916;
   Prof_PriceDA.Data[1098] := 0.1271916;
   Prof_PriceDA.Data[1099] := 0.1271916;
   Prof_PriceDA.Data[1100] := 0.1140588;
   Prof_PriceDA.Data[1101] := 0.1140588;
   Prof_PriceDA.Data[1102] := 0.1140588;
   Prof_PriceDA.Data[1103] := 0.1140588;
   Prof_PriceDA.Data[1104] := 0.1112292;
   Prof_PriceDA.Data[1105] := 0.1112292;
   Prof_PriceDA.Data[1106] := 0.1112292;
   Prof_PriceDA.Data[1107] := 0.1112292;
   Prof_PriceDA.Data[1108] := 0.1075788;
   Prof_PriceDA.Data[1109] := 0.1075788;
   Prof_PriceDA.Data[1110] := 0.1075788;
   Prof_PriceDA.Data[1111] := 0.1075788;
   Prof_PriceDA.Data[1112] := 0.1139616;
   Prof_PriceDA.Data[1113] := 0.1139616;
   Prof_PriceDA.Data[1114] := 0.1139616;
   Prof_PriceDA.Data[1115] := 0.1139616;
   Prof_PriceDA.Data[1116] := 0.1299564;
   Prof_PriceDA.Data[1117] := 0.1299564;
   Prof_PriceDA.Data[1118] := 0.1299564;
   Prof_PriceDA.Data[1119] := 0.1299564;
   Prof_PriceDA.Data[1120] := 0.1461024;
   Prof_PriceDA.Data[1121] := 0.1461024;
   Prof_PriceDA.Data[1122] := 0.1461024;
   Prof_PriceDA.Data[1123] := 0.1461024;
   Prof_PriceDA.Data[1124] := 0.1542564;
   Prof_PriceDA.Data[1125] := 0.1542564;
   Prof_PriceDA.Data[1126] := 0.1542564;
   Prof_PriceDA.Data[1127] := 0.1542564;
   Prof_PriceDA.Data[1128] := 0.1583928;
   Prof_PriceDA.Data[1129] := 0.1583928;
   Prof_PriceDA.Data[1130] := 0.1583928;
   Prof_PriceDA.Data[1131] := 0.1583928;
   Prof_PriceDA.Data[1132] := 0.1557468;
   Prof_PriceDA.Data[1133] := 0.1557468;
   Prof_PriceDA.Data[1134] := 0.1557468;
   Prof_PriceDA.Data[1135] := 0.1557468;
   Prof_PriceDA.Data[1136] := 0.1468152;
   Prof_PriceDA.Data[1137] := 0.1468152;
   Prof_PriceDA.Data[1138] := 0.1468152;
   Prof_PriceDA.Data[1139] := 0.1468152;
   Prof_PriceDA.Data[1140] := 0.1380348;
   Prof_PriceDA.Data[1141] := 0.1380348;
   Prof_PriceDA.Data[1142] := 0.1380348;
   Prof_PriceDA.Data[1143] := 0.1380348;
   Prof_PriceDA.Data[1144] := 0.1312956;
   Prof_PriceDA.Data[1145] := 0.1312956;
   Prof_PriceDA.Data[1146] := 0.1312956;
   Prof_PriceDA.Data[1147] := 0.1312956;
   Prof_PriceDA.Data[1148] := 0.124092;
   Prof_PriceDA.Data[1149] := 0.124092;
   Prof_PriceDA.Data[1150] := 0.124092;
   Prof_PriceDA.Data[1151] := 0.124092;
   Prof_PriceDA.Data[1152] := 0.1213812;
   Prof_PriceDA.Data[1153] := 0.1213812;
   Prof_PriceDA.Data[1154] := 0.1213812;
   Prof_PriceDA.Data[1155] := 0.1213812;
   Prof_PriceDA.Data[1156] := 0.1134756;
   Prof_PriceDA.Data[1157] := 0.1134756;
   Prof_PriceDA.Data[1158] := 0.1134756;
   Prof_PriceDA.Data[1159] := 0.1134756;
   Prof_PriceDA.Data[1160] := 0.1128168;
   Prof_PriceDA.Data[1161] := 0.1128168;
   Prof_PriceDA.Data[1162] := 0.1128168;
   Prof_PriceDA.Data[1163] := 0.1128168;
   Prof_PriceDA.Data[1164] := 0.1083996;
   Prof_PriceDA.Data[1165] := 0.1083996;
   Prof_PriceDA.Data[1166] := 0.1083996;
   Prof_PriceDA.Data[1167] := 0.1083996;
   Prof_PriceDA.Data[1168] := 0.108;
   Prof_PriceDA.Data[1169] := 0.108;
   Prof_PriceDA.Data[1170] := 0.108;
   Prof_PriceDA.Data[1171] := 0.108;
   Prof_PriceDA.Data[1172] := 0.1190052;
   Prof_PriceDA.Data[1173] := 0.1190052;
   Prof_PriceDA.Data[1174] := 0.1190052;
   Prof_PriceDA.Data[1175] := 0.1190052;
   Prof_PriceDA.Data[1176] := 0.1512108;
   Prof_PriceDA.Data[1177] := 0.1512108;
   Prof_PriceDA.Data[1178] := 0.1512108;
   Prof_PriceDA.Data[1179] := 0.1512108;
   Prof_PriceDA.Data[1180] := 0.1927476;
   Prof_PriceDA.Data[1181] := 0.1927476;
   Prof_PriceDA.Data[1182] := 0.1927476;
   Prof_PriceDA.Data[1183] := 0.1927476;
   Prof_PriceDA.Data[1184] := 0.2371032;
   Prof_PriceDA.Data[1185] := 0.2371032;
   Prof_PriceDA.Data[1186] := 0.2371032;
   Prof_PriceDA.Data[1187] := 0.2371032;
   Prof_PriceDA.Data[1188] := 0.1868184;
   Prof_PriceDA.Data[1189] := 0.1868184;
   Prof_PriceDA.Data[1190] := 0.1868184;
   Prof_PriceDA.Data[1191] := 0.1868184;
   Prof_PriceDA.Data[1192] := 0.15201;
   Prof_PriceDA.Data[1193] := 0.15201;
   Prof_PriceDA.Data[1194] := 0.15201;
   Prof_PriceDA.Data[1195] := 0.15201;
   Prof_PriceDA.Data[1196] := 0.1311444;
   Prof_PriceDA.Data[1197] := 0.1311444;
   Prof_PriceDA.Data[1198] := 0.1311444;
   Prof_PriceDA.Data[1199] := 0.1311444;
   Prof_PriceDA.Data[1200] := 0.1245456;
   Prof_PriceDA.Data[1201] := 0.1245456;
   Prof_PriceDA.Data[1202] := 0.1245456;
   Prof_PriceDA.Data[1203] := 0.1245456;
   Prof_PriceDA.Data[1204] := 0.1297512;
   Prof_PriceDA.Data[1205] := 0.1297512;
   Prof_PriceDA.Data[1206] := 0.1297512;
   Prof_PriceDA.Data[1207] := 0.1297512;
   Prof_PriceDA.Data[1208] := 0.1363284;
   Prof_PriceDA.Data[1209] := 0.1363284;
   Prof_PriceDA.Data[1210] := 0.1363284;
   Prof_PriceDA.Data[1211] := 0.1363284;
   Prof_PriceDA.Data[1212] := 0.1529928;
   Prof_PriceDA.Data[1213] := 0.1529928;
   Prof_PriceDA.Data[1214] := 0.1529928;
   Prof_PriceDA.Data[1215] := 0.1529928;
   Prof_PriceDA.Data[1216] := 0.1704564;
   Prof_PriceDA.Data[1217] := 0.1704564;
   Prof_PriceDA.Data[1218] := 0.1704564;
   Prof_PriceDA.Data[1219] := 0.1704564;
   Prof_PriceDA.Data[1220] := 0.1678212;
   Prof_PriceDA.Data[1221] := 0.1678212;
   Prof_PriceDA.Data[1222] := 0.1678212;
   Prof_PriceDA.Data[1223] := 0.1678212;
   Prof_PriceDA.Data[1224] := 0.16902;
   Prof_PriceDA.Data[1225] := 0.16902;
   Prof_PriceDA.Data[1226] := 0.16902;
   Prof_PriceDA.Data[1227] := 0.16902;
   Prof_PriceDA.Data[1228] := 0.1670976;
   Prof_PriceDA.Data[1229] := 0.1670976;
   Prof_PriceDA.Data[1230] := 0.1670976;
   Prof_PriceDA.Data[1231] := 0.1670976;
   Prof_PriceDA.Data[1232] := 0.1538244;
   Prof_PriceDA.Data[1233] := 0.1538244;
   Prof_PriceDA.Data[1234] := 0.1538244;
   Prof_PriceDA.Data[1235] := 0.1538244;
   Prof_PriceDA.Data[1236] := 0.1375164;
   Prof_PriceDA.Data[1237] := 0.1375164;
   Prof_PriceDA.Data[1238] := 0.1375164;
   Prof_PriceDA.Data[1239] := 0.1375164;
   Prof_PriceDA.Data[1240] := 0.1288008;
   Prof_PriceDA.Data[1241] := 0.1288008;
   Prof_PriceDA.Data[1242] := 0.1288008;
   Prof_PriceDA.Data[1243] := 0.1288008;
   Prof_PriceDA.Data[1244] := 0.1167588;
   Prof_PriceDA.Data[1245] := 0.1167588;
   Prof_PriceDA.Data[1246] := 0.1167588;
   Prof_PriceDA.Data[1247] := 0.1167588;
   Prof_PriceDA.Data[1248] := 0.1186812;
   Prof_PriceDA.Data[1249] := 0.1186812;
   Prof_PriceDA.Data[1250] := 0.1186812;
   Prof_PriceDA.Data[1251] := 0.1186812;
   Prof_PriceDA.Data[1252] := 0.115344;
   Prof_PriceDA.Data[1253] := 0.115344;
   Prof_PriceDA.Data[1254] := 0.115344;
   Prof_PriceDA.Data[1255] := 0.115344;
   Prof_PriceDA.Data[1256] := 0.1107;
   Prof_PriceDA.Data[1257] := 0.1107;
   Prof_PriceDA.Data[1258] := 0.1107;
   Prof_PriceDA.Data[1259] := 0.1107;
   Prof_PriceDA.Data[1260] := 0.1092312;
   Prof_PriceDA.Data[1261] := 0.1092312;
   Prof_PriceDA.Data[1262] := 0.1092312;
   Prof_PriceDA.Data[1263] := 0.1092312;
   Prof_PriceDA.Data[1264] := 0.1125036;
   Prof_PriceDA.Data[1265] := 0.1125036;
   Prof_PriceDA.Data[1266] := 0.1125036;
   Prof_PriceDA.Data[1267] := 0.1125036;
   Prof_PriceDA.Data[1268] := 0.1180332;
   Prof_PriceDA.Data[1269] := 0.1180332;
   Prof_PriceDA.Data[1270] := 0.1180332;
   Prof_PriceDA.Data[1271] := 0.1180332;
   Prof_PriceDA.Data[1272] := 0.1495908;
   Prof_PriceDA.Data[1273] := 0.1495908;
   Prof_PriceDA.Data[1274] := 0.1495908;
   Prof_PriceDA.Data[1275] := 0.1495908;
   Prof_PriceDA.Data[1276] := 0.1742688;
   Prof_PriceDA.Data[1277] := 0.1742688;
   Prof_PriceDA.Data[1278] := 0.1742688;
   Prof_PriceDA.Data[1279] := 0.1742688;
   Prof_PriceDA.Data[1280] := 0.2001672;
   Prof_PriceDA.Data[1281] := 0.2001672;
   Prof_PriceDA.Data[1282] := 0.2001672;
   Prof_PriceDA.Data[1283] := 0.2001672;
   Prof_PriceDA.Data[1284] := 0.16416;
   Prof_PriceDA.Data[1285] := 0.16416;
   Prof_PriceDA.Data[1286] := 0.16416;
   Prof_PriceDA.Data[1287] := 0.16416;
   Prof_PriceDA.Data[1288] := 0.141156;
   Prof_PriceDA.Data[1289] := 0.141156;
   Prof_PriceDA.Data[1290] := 0.141156;
   Prof_PriceDA.Data[1291] := 0.141156;
   Prof_PriceDA.Data[1292] := 0.1340712;
   Prof_PriceDA.Data[1293] := 0.1340712;
   Prof_PriceDA.Data[1294] := 0.1340712;
   Prof_PriceDA.Data[1295] := 0.1340712;
   Prof_PriceDA.Data[1296] := 0.1289304;
   Prof_PriceDA.Data[1297] := 0.1289304;
   Prof_PriceDA.Data[1298] := 0.1289304;
   Prof_PriceDA.Data[1299] := 0.1289304;
   Prof_PriceDA.Data[1300] := 0.1293084;
   Prof_PriceDA.Data[1301] := 0.1293084;
   Prof_PriceDA.Data[1302] := 0.1293084;
   Prof_PriceDA.Data[1303] := 0.1293084;
   Prof_PriceDA.Data[1304] := 0.1439532;
   Prof_PriceDA.Data[1305] := 0.1439532;
   Prof_PriceDA.Data[1306] := 0.1439532;
   Prof_PriceDA.Data[1307] := 0.1439532;
   Prof_PriceDA.Data[1308] := 0.1770552;
   Prof_PriceDA.Data[1309] := 0.1770552;
   Prof_PriceDA.Data[1310] := 0.1770552;
   Prof_PriceDA.Data[1311] := 0.1770552;
   Prof_PriceDA.Data[1312] := 0.1979964;
   Prof_PriceDA.Data[1313] := 0.1979964;
   Prof_PriceDA.Data[1314] := 0.1979964;
   Prof_PriceDA.Data[1315] := 0.1979964;
   Prof_PriceDA.Data[1316] := 0.2446632;
   Prof_PriceDA.Data[1317] := 0.2446632;
   Prof_PriceDA.Data[1318] := 0.2446632;
   Prof_PriceDA.Data[1319] := 0.2446632;
   Prof_PriceDA.Data[1320] := 0.239652;
   Prof_PriceDA.Data[1321] := 0.239652;
   Prof_PriceDA.Data[1322] := 0.239652;
   Prof_PriceDA.Data[1323] := 0.239652;
   Prof_PriceDA.Data[1324] := 0.211572;
   Prof_PriceDA.Data[1325] := 0.211572;
   Prof_PriceDA.Data[1326] := 0.211572;
   Prof_PriceDA.Data[1327] := 0.211572;
   Prof_PriceDA.Data[1328] := 0.187164;
   Prof_PriceDA.Data[1329] := 0.187164;
   Prof_PriceDA.Data[1330] := 0.187164;
   Prof_PriceDA.Data[1331] := 0.187164;
   Prof_PriceDA.Data[1332] := 0.172746;
   Prof_PriceDA.Data[1333] := 0.172746;
   Prof_PriceDA.Data[1334] := 0.172746;
   Prof_PriceDA.Data[1335] := 0.172746;
   Prof_PriceDA.Data[1336] := 0.1610172;
   Prof_PriceDA.Data[1337] := 0.1610172;
   Prof_PriceDA.Data[1338] := 0.1610172;
   Prof_PriceDA.Data[1339] := 0.1610172;
   Prof_PriceDA.Data[1340] := 0.1348812;
   Prof_PriceDA.Data[1341] := 0.1348812;
   Prof_PriceDA.Data[1342] := 0.1348812;
   Prof_PriceDA.Data[1343] := 0.1348812;
   Prof_PriceDA.Data[1344] := 0.127656;
   Prof_PriceDA.Data[1345] := 0.127656;
   Prof_PriceDA.Data[1346] := 0.127656;
   Prof_PriceDA.Data[1347] := 0.127656;
   Prof_PriceDA.Data[1348] := 0.1213488;
   Prof_PriceDA.Data[1349] := 0.1213488;
   Prof_PriceDA.Data[1350] := 0.1213488;
   Prof_PriceDA.Data[1351] := 0.1213488;
   Prof_PriceDA.Data[1352] := 0.1200528;
   Prof_PriceDA.Data[1353] := 0.1200528;
   Prof_PriceDA.Data[1354] := 0.1200528;
   Prof_PriceDA.Data[1355] := 0.1200528;
   Prof_PriceDA.Data[1356] := 0.1174932;
   Prof_PriceDA.Data[1357] := 0.1174932;
   Prof_PriceDA.Data[1358] := 0.1174932;
   Prof_PriceDA.Data[1359] := 0.1174932;
   Prof_PriceDA.Data[1360] := 0.1255068;
   Prof_PriceDA.Data[1361] := 0.1255068;
   Prof_PriceDA.Data[1362] := 0.1255068;
   Prof_PriceDA.Data[1363] := 0.1255068;
   Prof_PriceDA.Data[1364] := 0.1390392;
   Prof_PriceDA.Data[1365] := 0.1390392;
   Prof_PriceDA.Data[1366] := 0.1390392;
   Prof_PriceDA.Data[1367] := 0.1390392;
   Prof_PriceDA.Data[1368] := 0.1600992;
   Prof_PriceDA.Data[1369] := 0.1600992;
   Prof_PriceDA.Data[1370] := 0.1600992;
   Prof_PriceDA.Data[1371] := 0.1600992;
   Prof_PriceDA.Data[1372] := 0.2120148;
   Prof_PriceDA.Data[1373] := 0.2120148;
   Prof_PriceDA.Data[1374] := 0.2120148;
   Prof_PriceDA.Data[1375] := 0.2120148;
   Prof_PriceDA.Data[1376] := 0.3359124;
   Prof_PriceDA.Data[1377] := 0.3359124;
   Prof_PriceDA.Data[1378] := 0.3359124;
   Prof_PriceDA.Data[1379] := 0.3359124;
   Prof_PriceDA.Data[1380] := 0.338904;
   Prof_PriceDA.Data[1381] := 0.338904;
   Prof_PriceDA.Data[1382] := 0.338904;
   Prof_PriceDA.Data[1383] := 0.338904;
   Prof_PriceDA.Data[1384] := 0.3266568;
   Prof_PriceDA.Data[1385] := 0.3266568;
   Prof_PriceDA.Data[1386] := 0.3266568;
   Prof_PriceDA.Data[1387] := 0.3266568;
   Prof_PriceDA.Data[1388] := 0.325566;
   Prof_PriceDA.Data[1389] := 0.325566;
   Prof_PriceDA.Data[1390] := 0.325566;
   Prof_PriceDA.Data[1391] := 0.325566;
   Prof_PriceDA.Data[1392] := 0.31023;
   Prof_PriceDA.Data[1393] := 0.31023;
   Prof_PriceDA.Data[1394] := 0.31023;
   Prof_PriceDA.Data[1395] := 0.31023;
   Prof_PriceDA.Data[1396] := 0.306774;
   Prof_PriceDA.Data[1397] := 0.306774;
   Prof_PriceDA.Data[1398] := 0.306774;
   Prof_PriceDA.Data[1399] := 0.306774;
   Prof_PriceDA.Data[1400] := 0.3062448;
   Prof_PriceDA.Data[1401] := 0.3062448;
   Prof_PriceDA.Data[1402] := 0.3062448;
   Prof_PriceDA.Data[1403] := 0.3062448;
   Prof_PriceDA.Data[1404] := 0.3319596;
   Prof_PriceDA.Data[1405] := 0.3319596;
   Prof_PriceDA.Data[1406] := 0.3319596;
   Prof_PriceDA.Data[1407] := 0.3319596;
   Prof_PriceDA.Data[1408] := 0.326268;
   Prof_PriceDA.Data[1409] := 0.326268;
   Prof_PriceDA.Data[1410] := 0.326268;
   Prof_PriceDA.Data[1411] := 0.326268;
   Prof_PriceDA.Data[1412] := 0.368226;
   Prof_PriceDA.Data[1413] := 0.368226;
   Prof_PriceDA.Data[1414] := 0.368226;
   Prof_PriceDA.Data[1415] := 0.368226;
   Prof_PriceDA.Data[1416] := 0.320328;
   Prof_PriceDA.Data[1417] := 0.320328;
   Prof_PriceDA.Data[1418] := 0.320328;
   Prof_PriceDA.Data[1419] := 0.320328;
   Prof_PriceDA.Data[1420] := 0.265248;
   Prof_PriceDA.Data[1421] := 0.265248;
   Prof_PriceDA.Data[1422] := 0.265248;
   Prof_PriceDA.Data[1423] := 0.265248;
   Prof_PriceDA.Data[1424] := 0.1937088;
   Prof_PriceDA.Data[1425] := 0.1937088;
   Prof_PriceDA.Data[1426] := 0.1937088;
   Prof_PriceDA.Data[1427] := 0.1937088;
   Prof_PriceDA.Data[1428] := 0.1670328;
   Prof_PriceDA.Data[1429] := 0.1670328;
   Prof_PriceDA.Data[1430] := 0.1670328;
   Prof_PriceDA.Data[1431] := 0.1670328;
   Prof_PriceDA.Data[1432] := 0.1554768;
   Prof_PriceDA.Data[1433] := 0.1554768;
   Prof_PriceDA.Data[1434] := 0.1554768;
   Prof_PriceDA.Data[1435] := 0.1554768;
   Prof_PriceDA.Data[1436] := 0.133812;
   Prof_PriceDA.Data[1437] := 0.133812;
   Prof_PriceDA.Data[1438] := 0.133812;
   Prof_PriceDA.Data[1439] := 0.133812;
   Prof_PriceDA.Data[1440] := 0.136296;
   Prof_PriceDA.Data[1441] := 0.136296;
   Prof_PriceDA.Data[1442] := 0.136296;
   Prof_PriceDA.Data[1443] := 0.136296;
   Prof_PriceDA.Data[1444] := 0.131868;
   Prof_PriceDA.Data[1445] := 0.131868;
   Prof_PriceDA.Data[1446] := 0.131868;
   Prof_PriceDA.Data[1447] := 0.131868;
   Prof_PriceDA.Data[1448] := 0.1281636;
   Prof_PriceDA.Data[1449] := 0.1281636;
   Prof_PriceDA.Data[1450] := 0.1281636;
   Prof_PriceDA.Data[1451] := 0.1281636;
   Prof_PriceDA.Data[1452] := 0.1259928;
   Prof_PriceDA.Data[1453] := 0.1259928;
   Prof_PriceDA.Data[1454] := 0.1259928;
   Prof_PriceDA.Data[1455] := 0.1259928;
   Prof_PriceDA.Data[1456] := 0.1292652;
   Prof_PriceDA.Data[1457] := 0.1292652;
   Prof_PriceDA.Data[1458] := 0.1292652;
   Prof_PriceDA.Data[1459] := 0.1292652;
   Prof_PriceDA.Data[1460] := 0.1392012;
   Prof_PriceDA.Data[1461] := 0.1392012;
   Prof_PriceDA.Data[1462] := 0.1392012;
   Prof_PriceDA.Data[1463] := 0.1392012;
   Prof_PriceDA.Data[1464] := 0.1701216;
   Prof_PriceDA.Data[1465] := 0.1701216;
   Prof_PriceDA.Data[1466] := 0.1701216;
   Prof_PriceDA.Data[1467] := 0.1701216;
   Prof_PriceDA.Data[1468] := 0.2121984;
   Prof_PriceDA.Data[1469] := 0.2121984;
   Prof_PriceDA.Data[1470] := 0.2121984;
   Prof_PriceDA.Data[1471] := 0.2121984;
   Prof_PriceDA.Data[1472] := 0.2210544;
   Prof_PriceDA.Data[1473] := 0.2210544;
   Prof_PriceDA.Data[1474] := 0.2210544;
   Prof_PriceDA.Data[1475] := 0.2210544;
   Prof_PriceDA.Data[1476] := 0.189;
   Prof_PriceDA.Data[1477] := 0.189;
   Prof_PriceDA.Data[1478] := 0.189;
   Prof_PriceDA.Data[1479] := 0.189;
   Prof_PriceDA.Data[1480] := 0.164052;
   Prof_PriceDA.Data[1481] := 0.164052;
   Prof_PriceDA.Data[1482] := 0.164052;
   Prof_PriceDA.Data[1483] := 0.164052;
   Prof_PriceDA.Data[1484] := 0.1518912;
   Prof_PriceDA.Data[1485] := 0.1518912;
   Prof_PriceDA.Data[1486] := 0.1518912;
   Prof_PriceDA.Data[1487] := 0.1518912;
   Prof_PriceDA.Data[1488] := 0.1456488;
   Prof_PriceDA.Data[1489] := 0.1456488;
   Prof_PriceDA.Data[1490] := 0.1456488;
   Prof_PriceDA.Data[1491] := 0.1456488;
   Prof_PriceDA.Data[1492] := 0.1492344;
   Prof_PriceDA.Data[1493] := 0.1492344;
   Prof_PriceDA.Data[1494] := 0.1492344;
   Prof_PriceDA.Data[1495] := 0.1492344;
   Prof_PriceDA.Data[1496] := 0.1566;
   Prof_PriceDA.Data[1497] := 0.1566;
   Prof_PriceDA.Data[1498] := 0.1566;
   Prof_PriceDA.Data[1499] := 0.1566;
   Prof_PriceDA.Data[1500] := 0.1827144;
   Prof_PriceDA.Data[1501] := 0.1827144;
   Prof_PriceDA.Data[1502] := 0.1827144;
   Prof_PriceDA.Data[1503] := 0.1827144;
   Prof_PriceDA.Data[1504] := 0.19683;
   Prof_PriceDA.Data[1505] := 0.19683;
   Prof_PriceDA.Data[1506] := 0.19683;
   Prof_PriceDA.Data[1507] := 0.19683;
   Prof_PriceDA.Data[1508] := 0.2082348;
   Prof_PriceDA.Data[1509] := 0.2082348;
   Prof_PriceDA.Data[1510] := 0.2082348;
   Prof_PriceDA.Data[1511] := 0.2082348;
   Prof_PriceDA.Data[1512] := 0.1990656;
   Prof_PriceDA.Data[1513] := 0.1990656;
   Prof_PriceDA.Data[1514] := 0.1990656;
   Prof_PriceDA.Data[1515] := 0.1990656;
   Prof_PriceDA.Data[1516] := 0.1943676;
   Prof_PriceDA.Data[1517] := 0.1943676;
   Prof_PriceDA.Data[1518] := 0.1943676;
   Prof_PriceDA.Data[1519] := 0.1943676;
   Prof_PriceDA.Data[1520] := 0.172368;
   Prof_PriceDA.Data[1521] := 0.172368;
   Prof_PriceDA.Data[1522] := 0.172368;
   Prof_PriceDA.Data[1523] := 0.172368;
   Prof_PriceDA.Data[1524] := 0.1623996;
   Prof_PriceDA.Data[1525] := 0.1623996;
   Prof_PriceDA.Data[1526] := 0.1623996;
   Prof_PriceDA.Data[1527] := 0.1623996;
   Prof_PriceDA.Data[1528] := 0.1519992;
   Prof_PriceDA.Data[1529] := 0.1519992;
   Prof_PriceDA.Data[1530] := 0.1519992;
   Prof_PriceDA.Data[1531] := 0.1519992;
   Prof_PriceDA.Data[1532] := 0.1398276;
   Prof_PriceDA.Data[1533] := 0.1398276;
   Prof_PriceDA.Data[1534] := 0.1398276;
   Prof_PriceDA.Data[1535] := 0.1398276;
   Prof_PriceDA.Data[1536] := 0.1364364;
   Prof_PriceDA.Data[1537] := 0.1364364;
   Prof_PriceDA.Data[1538] := 0.1364364;
   Prof_PriceDA.Data[1539] := 0.1364364;
   Prof_PriceDA.Data[1540] := 0.1331208;
   Prof_PriceDA.Data[1541] := 0.1331208;
   Prof_PriceDA.Data[1542] := 0.1331208;
   Prof_PriceDA.Data[1543] := 0.1331208;
   Prof_PriceDA.Data[1544] := 0.1297836;
   Prof_PriceDA.Data[1545] := 0.1297836;
   Prof_PriceDA.Data[1546] := 0.1297836;
   Prof_PriceDA.Data[1547] := 0.1297836;
   Prof_PriceDA.Data[1548] := 0.1277532;
   Prof_PriceDA.Data[1549] := 0.1277532;
   Prof_PriceDA.Data[1550] := 0.1277532;
   Prof_PriceDA.Data[1551] := 0.1277532;
   Prof_PriceDA.Data[1552] := 0.1277964;
   Prof_PriceDA.Data[1553] := 0.1277964;
   Prof_PriceDA.Data[1554] := 0.1277964;
   Prof_PriceDA.Data[1555] := 0.1277964;
   Prof_PriceDA.Data[1556] := 0.1346328;
   Prof_PriceDA.Data[1557] := 0.1346328;
   Prof_PriceDA.Data[1558] := 0.1346328;
   Prof_PriceDA.Data[1559] := 0.1346328;
   Prof_PriceDA.Data[1560] := 0.152064;
   Prof_PriceDA.Data[1561] := 0.152064;
   Prof_PriceDA.Data[1562] := 0.152064;
   Prof_PriceDA.Data[1563] := 0.152064;
   Prof_PriceDA.Data[1564] := 0.1890108;
   Prof_PriceDA.Data[1565] := 0.1890108;
   Prof_PriceDA.Data[1566] := 0.1890108;
   Prof_PriceDA.Data[1567] := 0.1890108;
   Prof_PriceDA.Data[1568] := 0.2247804;
   Prof_PriceDA.Data[1569] := 0.2247804;
   Prof_PriceDA.Data[1570] := 0.2247804;
   Prof_PriceDA.Data[1571] := 0.2247804;
   Prof_PriceDA.Data[1572] := 0.1893672;
   Prof_PriceDA.Data[1573] := 0.1893672;
   Prof_PriceDA.Data[1574] := 0.1893672;
   Prof_PriceDA.Data[1575] := 0.1893672;
   Prof_PriceDA.Data[1576] := 0.1700352;
   Prof_PriceDA.Data[1577] := 0.1700352;
   Prof_PriceDA.Data[1578] := 0.1700352;
   Prof_PriceDA.Data[1579] := 0.1700352;
   Prof_PriceDA.Data[1580] := 0.1518696;
   Prof_PriceDA.Data[1581] := 0.1518696;
   Prof_PriceDA.Data[1582] := 0.1518696;
   Prof_PriceDA.Data[1583] := 0.1518696;
   Prof_PriceDA.Data[1584] := 0.1365552;
   Prof_PriceDA.Data[1585] := 0.1365552;
   Prof_PriceDA.Data[1586] := 0.1365552;
   Prof_PriceDA.Data[1587] := 0.1365552;
   Prof_PriceDA.Data[1588] := 0.1339524;
   Prof_PriceDA.Data[1589] := 0.1339524;
   Prof_PriceDA.Data[1590] := 0.1339524;
   Prof_PriceDA.Data[1591] := 0.1339524;
   Prof_PriceDA.Data[1592] := 0.1444284;
   Prof_PriceDA.Data[1593] := 0.1444284;
   Prof_PriceDA.Data[1594] := 0.1444284;
   Prof_PriceDA.Data[1595] := 0.1444284;
   Prof_PriceDA.Data[1596] := 0.1637172;
   Prof_PriceDA.Data[1597] := 0.1637172;
   Prof_PriceDA.Data[1598] := 0.1637172;
   Prof_PriceDA.Data[1599] := 0.1637172;
   Prof_PriceDA.Data[1600] := 0.1839888;
   Prof_PriceDA.Data[1601] := 0.1839888;
   Prof_PriceDA.Data[1602] := 0.1839888;
   Prof_PriceDA.Data[1603] := 0.1839888;
   Prof_PriceDA.Data[1604] := 0.1930284;
   Prof_PriceDA.Data[1605] := 0.1930284;
   Prof_PriceDA.Data[1606] := 0.1930284;
   Prof_PriceDA.Data[1607] := 0.1930284;
   Prof_PriceDA.Data[1608] := 0.1943136;
   Prof_PriceDA.Data[1609] := 0.1943136;
   Prof_PriceDA.Data[1610] := 0.1943136;
   Prof_PriceDA.Data[1611] := 0.1943136;
   Prof_PriceDA.Data[1612] := 0.1881576;
   Prof_PriceDA.Data[1613] := 0.1881576;
   Prof_PriceDA.Data[1614] := 0.1881576;
   Prof_PriceDA.Data[1615] := 0.1881576;
   Prof_PriceDA.Data[1616] := 0.1705428;
   Prof_PriceDA.Data[1617] := 0.1705428;
   Prof_PriceDA.Data[1618] := 0.1705428;
   Prof_PriceDA.Data[1619] := 0.1705428;
   Prof_PriceDA.Data[1620] := 0.1566;
   Prof_PriceDA.Data[1621] := 0.1566;
   Prof_PriceDA.Data[1622] := 0.1566;
   Prof_PriceDA.Data[1623] := 0.1566;
   Prof_PriceDA.Data[1624] := 0.1511676;
   Prof_PriceDA.Data[1625] := 0.1511676;
   Prof_PriceDA.Data[1626] := 0.1511676;
   Prof_PriceDA.Data[1627] := 0.1511676;
   Prof_PriceDA.Data[1628] := 0.1383588;
   Prof_PriceDA.Data[1629] := 0.1383588;
   Prof_PriceDA.Data[1630] := 0.1383588;
   Prof_PriceDA.Data[1631] := 0.1383588;
   Prof_PriceDA.Data[1632] := 0.1363392;
   Prof_PriceDA.Data[1633] := 0.1363392;
   Prof_PriceDA.Data[1634] := 0.1363392;
   Prof_PriceDA.Data[1635] := 0.1363392;
   Prof_PriceDA.Data[1636] := 0.1309284;
   Prof_PriceDA.Data[1637] := 0.1309284;
   Prof_PriceDA.Data[1638] := 0.1309284;
   Prof_PriceDA.Data[1639] := 0.1309284;
   Prof_PriceDA.Data[1640] := 0.1311336;
   Prof_PriceDA.Data[1641] := 0.1311336;
   Prof_PriceDA.Data[1642] := 0.1311336;
   Prof_PriceDA.Data[1643] := 0.1311336;
   Prof_PriceDA.Data[1644] := 0.128412;
   Prof_PriceDA.Data[1645] := 0.128412;
   Prof_PriceDA.Data[1646] := 0.128412;
   Prof_PriceDA.Data[1647] := 0.128412;
   Prof_PriceDA.Data[1648] := 0.1263816;
   Prof_PriceDA.Data[1649] := 0.1263816;
   Prof_PriceDA.Data[1650] := 0.1263816;
   Prof_PriceDA.Data[1651] := 0.1263816;
   Prof_PriceDA.Data[1652] := 0.1294164;
   Prof_PriceDA.Data[1653] := 0.1294164;
   Prof_PriceDA.Data[1654] := 0.1294164;
   Prof_PriceDA.Data[1655] := 0.1294164;
   Prof_PriceDA.Data[1656] := 0.1325592;
   Prof_PriceDA.Data[1657] := 0.1325592;
   Prof_PriceDA.Data[1658] := 0.1325592;
   Prof_PriceDA.Data[1659] := 0.1325592;
   Prof_PriceDA.Data[1660] := 0.1465776;
   Prof_PriceDA.Data[1661] := 0.1465776;
   Prof_PriceDA.Data[1662] := 0.1465776;
   Prof_PriceDA.Data[1663] := 0.1465776;
   Prof_PriceDA.Data[1664] := 0.157626;
   Prof_PriceDA.Data[1665] := 0.157626;
   Prof_PriceDA.Data[1666] := 0.157626;
   Prof_PriceDA.Data[1667] := 0.157626;
   Prof_PriceDA.Data[1668] := 0.155628;
   Prof_PriceDA.Data[1669] := 0.155628;
   Prof_PriceDA.Data[1670] := 0.155628;
   Prof_PriceDA.Data[1671] := 0.155628;
   Prof_PriceDA.Data[1672] := 0.1445796;
   Prof_PriceDA.Data[1673] := 0.1445796;
   Prof_PriceDA.Data[1674] := 0.1445796;
   Prof_PriceDA.Data[1675] := 0.1445796;
   Prof_PriceDA.Data[1676] := 0.1315224;
   Prof_PriceDA.Data[1677] := 0.1315224;
   Prof_PriceDA.Data[1678] := 0.1315224;
   Prof_PriceDA.Data[1679] := 0.1315224;
   Prof_PriceDA.Data[1680] := 0.1283796;
   Prof_PriceDA.Data[1681] := 0.1283796;
   Prof_PriceDA.Data[1682] := 0.1283796;
   Prof_PriceDA.Data[1683] := 0.1283796;
   Prof_PriceDA.Data[1684] := 0.1242108;
   Prof_PriceDA.Data[1685] := 0.1242108;
   Prof_PriceDA.Data[1686] := 0.1242108;
   Prof_PriceDA.Data[1687] := 0.1242108;
   Prof_PriceDA.Data[1688] := 0.129168;
   Prof_PriceDA.Data[1689] := 0.129168;
   Prof_PriceDA.Data[1690] := 0.129168;
   Prof_PriceDA.Data[1691] := 0.129168;
   Prof_PriceDA.Data[1692] := 0.149094;
   Prof_PriceDA.Data[1693] := 0.149094;
   Prof_PriceDA.Data[1694] := 0.149094;
   Prof_PriceDA.Data[1695] := 0.149094;
   Prof_PriceDA.Data[1696] := 0.1772712;
   Prof_PriceDA.Data[1697] := 0.1772712;
   Prof_PriceDA.Data[1698] := 0.1772712;
   Prof_PriceDA.Data[1699] := 0.1772712;
   Prof_PriceDA.Data[1700] := 0.1826928;
   Prof_PriceDA.Data[1701] := 0.1826928;
   Prof_PriceDA.Data[1702] := 0.1826928;
   Prof_PriceDA.Data[1703] := 0.1826928;
   Prof_PriceDA.Data[1704] := 0.1809756;
   Prof_PriceDA.Data[1705] := 0.1809756;
   Prof_PriceDA.Data[1706] := 0.1809756;
   Prof_PriceDA.Data[1707] := 0.1809756;
   Prof_PriceDA.Data[1708] := 0.181278;
   Prof_PriceDA.Data[1709] := 0.181278;
   Prof_PriceDA.Data[1710] := 0.181278;
   Prof_PriceDA.Data[1711] := 0.181278;
   Prof_PriceDA.Data[1712] := 0.1686096;
   Prof_PriceDA.Data[1713] := 0.1686096;
   Prof_PriceDA.Data[1714] := 0.1686096;
   Prof_PriceDA.Data[1715] := 0.1686096;
   Prof_PriceDA.Data[1716] := 0.1548936;
   Prof_PriceDA.Data[1717] := 0.1548936;
   Prof_PriceDA.Data[1718] := 0.1548936;
   Prof_PriceDA.Data[1719] := 0.1548936;
   Prof_PriceDA.Data[1720] := 0.147312;
   Prof_PriceDA.Data[1721] := 0.147312;
   Prof_PriceDA.Data[1722] := 0.147312;
   Prof_PriceDA.Data[1723] := 0.147312;
   Prof_PriceDA.Data[1724] := 0.1397088;
   Prof_PriceDA.Data[1725] := 0.1397088;
   Prof_PriceDA.Data[1726] := 0.1397088;
   Prof_PriceDA.Data[1727] := 0.1397088;
   Prof_PriceDA.Data[1728] := 0.1403028;
   Prof_PriceDA.Data[1729] := 0.1403028;
   Prof_PriceDA.Data[1730] := 0.1403028;
   Prof_PriceDA.Data[1731] := 0.1403028;
   Prof_PriceDA.Data[1732] := 0.1350108;
   Prof_PriceDA.Data[1733] := 0.1350108;
   Prof_PriceDA.Data[1734] := 0.1350108;
   Prof_PriceDA.Data[1735] := 0.1350108;
   Prof_PriceDA.Data[1736] := 0.1336068;
   Prof_PriceDA.Data[1737] := 0.1336068;
   Prof_PriceDA.Data[1738] := 0.1336068;
   Prof_PriceDA.Data[1739] := 0.1336068;
   Prof_PriceDA.Data[1740] := 0.1309392;
   Prof_PriceDA.Data[1741] := 0.1309392;
   Prof_PriceDA.Data[1742] := 0.1309392;
   Prof_PriceDA.Data[1743] := 0.1309392;
   Prof_PriceDA.Data[1744] := 0.1297944;
   Prof_PriceDA.Data[1745] := 0.1297944;
   Prof_PriceDA.Data[1746] := 0.1297944;
   Prof_PriceDA.Data[1747] := 0.1297944;
   Prof_PriceDA.Data[1748] := 0.1296;
   Prof_PriceDA.Data[1749] := 0.1296;
   Prof_PriceDA.Data[1750] := 0.1296;
   Prof_PriceDA.Data[1751] := 0.1296;
   Prof_PriceDA.Data[1752] := 0.1314252;
   Prof_PriceDA.Data[1753] := 0.1314252;
   Prof_PriceDA.Data[1754] := 0.1314252;
   Prof_PriceDA.Data[1755] := 0.1314252;
   Prof_PriceDA.Data[1756] := 0.1340172;
   Prof_PriceDA.Data[1757] := 0.1340172;
   Prof_PriceDA.Data[1758] := 0.1340172;
   Prof_PriceDA.Data[1759] := 0.1340172;
   Prof_PriceDA.Data[1760] := 0.1335636;
   Prof_PriceDA.Data[1761] := 0.1335636;
   Prof_PriceDA.Data[1762] := 0.1335636;
   Prof_PriceDA.Data[1763] := 0.1335636;
   Prof_PriceDA.Data[1764] := 0.136188;
   Prof_PriceDA.Data[1765] := 0.136188;
   Prof_PriceDA.Data[1766] := 0.136188;
   Prof_PriceDA.Data[1767] := 0.136188;
   Prof_PriceDA.Data[1768] := 0.1366092;
   Prof_PriceDA.Data[1769] := 0.1366092;
   Prof_PriceDA.Data[1770] := 0.1366092;
   Prof_PriceDA.Data[1771] := 0.1366092;
   Prof_PriceDA.Data[1772] := 0.1341252;
   Prof_PriceDA.Data[1773] := 0.1341252;
   Prof_PriceDA.Data[1774] := 0.1341252;
   Prof_PriceDA.Data[1775] := 0.1341252;
   Prof_PriceDA.Data[1776] := 0.12123;
   Prof_PriceDA.Data[1777] := 0.12123;
   Prof_PriceDA.Data[1778] := 0.12123;
   Prof_PriceDA.Data[1779] := 0.12123;
   Prof_PriceDA.Data[1780] := 0.1161108;
   Prof_PriceDA.Data[1781] := 0.1161108;
   Prof_PriceDA.Data[1782] := 0.1161108;
   Prof_PriceDA.Data[1783] := 0.1161108;
   Prof_PriceDA.Data[1784] := 0.1261548;
   Prof_PriceDA.Data[1785] := 0.1261548;
   Prof_PriceDA.Data[1786] := 0.1261548;
   Prof_PriceDA.Data[1787] := 0.1261548;
   Prof_PriceDA.Data[1788] := 0.1377324;
   Prof_PriceDA.Data[1789] := 0.1377324;
   Prof_PriceDA.Data[1790] := 0.1377324;
   Prof_PriceDA.Data[1791] := 0.1377324;
   Prof_PriceDA.Data[1792] := 0.1627344;
   Prof_PriceDA.Data[1793] := 0.1627344;
   Prof_PriceDA.Data[1794] := 0.1627344;
   Prof_PriceDA.Data[1795] := 0.1627344;
   Prof_PriceDA.Data[1796] := 0.1759428;
   Prof_PriceDA.Data[1797] := 0.1759428;
   Prof_PriceDA.Data[1798] := 0.1759428;
   Prof_PriceDA.Data[1799] := 0.1759428;
   Prof_PriceDA.Data[1800] := 0.180522;
   Prof_PriceDA.Data[1801] := 0.180522;
   Prof_PriceDA.Data[1802] := 0.180522;
   Prof_PriceDA.Data[1803] := 0.180522;
   Prof_PriceDA.Data[1804] := 0.1794096;
   Prof_PriceDA.Data[1805] := 0.1794096;
   Prof_PriceDA.Data[1806] := 0.1794096;
   Prof_PriceDA.Data[1807] := 0.1794096;
   Prof_PriceDA.Data[1808] := 0.1741608;
   Prof_PriceDA.Data[1809] := 0.1741608;
   Prof_PriceDA.Data[1810] := 0.1741608;
   Prof_PriceDA.Data[1811] := 0.1741608;
   Prof_PriceDA.Data[1812] := 0.1651644;
   Prof_PriceDA.Data[1813] := 0.1651644;
   Prof_PriceDA.Data[1814] := 0.1651644;
   Prof_PriceDA.Data[1815] := 0.1651644;
   Prof_PriceDA.Data[1816] := 0.145044;
   Prof_PriceDA.Data[1817] := 0.145044;
   Prof_PriceDA.Data[1818] := 0.145044;
   Prof_PriceDA.Data[1819] := 0.145044;
   Prof_PriceDA.Data[1820] := 0.133866;
   Prof_PriceDA.Data[1821] := 0.133866;
   Prof_PriceDA.Data[1822] := 0.133866;
   Prof_PriceDA.Data[1823] := 0.133866;
   Prof_PriceDA.Data[1824] := 0.1322784;
   Prof_PriceDA.Data[1825] := 0.1322784;
   Prof_PriceDA.Data[1826] := 0.1322784;
   Prof_PriceDA.Data[1827] := 0.1322784;
   Prof_PriceDA.Data[1828] := 0.1294056;
   Prof_PriceDA.Data[1829] := 0.1294056;
   Prof_PriceDA.Data[1830] := 0.1294056;
   Prof_PriceDA.Data[1831] := 0.1294056;
   Prof_PriceDA.Data[1832] := 0.1259388;
   Prof_PriceDA.Data[1833] := 0.1259388;
   Prof_PriceDA.Data[1834] := 0.1259388;
   Prof_PriceDA.Data[1835] := 0.1259388;
   Prof_PriceDA.Data[1836] := 0.1235628;
   Prof_PriceDA.Data[1837] := 0.1235628;
   Prof_PriceDA.Data[1838] := 0.1235628;
   Prof_PriceDA.Data[1839] := 0.1235628;
   Prof_PriceDA.Data[1840] := 0.124686;
   Prof_PriceDA.Data[1841] := 0.124686;
   Prof_PriceDA.Data[1842] := 0.124686;
   Prof_PriceDA.Data[1843] := 0.124686;
   Prof_PriceDA.Data[1844] := 0.1404216;
   Prof_PriceDA.Data[1845] := 0.1404216;
   Prof_PriceDA.Data[1846] := 0.1404216;
   Prof_PriceDA.Data[1847] := 0.1404216;
   Prof_PriceDA.Data[1848] := 0.1766232;
   Prof_PriceDA.Data[1849] := 0.1766232;
   Prof_PriceDA.Data[1850] := 0.1766232;
   Prof_PriceDA.Data[1851] := 0.1766232;
   Prof_PriceDA.Data[1852] := 0.3070548;
   Prof_PriceDA.Data[1853] := 0.3070548;
   Prof_PriceDA.Data[1854] := 0.3070548;
   Prof_PriceDA.Data[1855] := 0.3070548;
   Prof_PriceDA.Data[1856] := 0.4670028;
   Prof_PriceDA.Data[1857] := 0.4670028;
   Prof_PriceDA.Data[1858] := 0.4670028;
   Prof_PriceDA.Data[1859] := 0.4670028;
   Prof_PriceDA.Data[1860] := 0.3149496;
   Prof_PriceDA.Data[1861] := 0.3149496;
   Prof_PriceDA.Data[1862] := 0.3149496;
   Prof_PriceDA.Data[1863] := 0.3149496;
   Prof_PriceDA.Data[1864] := 0.2551932;
   Prof_PriceDA.Data[1865] := 0.2551932;
   Prof_PriceDA.Data[1866] := 0.2551932;
   Prof_PriceDA.Data[1867] := 0.2551932;
   Prof_PriceDA.Data[1868] := 0.2076084;
   Prof_PriceDA.Data[1869] := 0.2076084;
   Prof_PriceDA.Data[1870] := 0.2076084;
   Prof_PriceDA.Data[1871] := 0.2076084;
   Prof_PriceDA.Data[1872] := 0.193266;
   Prof_PriceDA.Data[1873] := 0.193266;
   Prof_PriceDA.Data[1874] := 0.193266;
   Prof_PriceDA.Data[1875] := 0.193266;
   Prof_PriceDA.Data[1876] := 0.1851012;
   Prof_PriceDA.Data[1877] := 0.1851012;
   Prof_PriceDA.Data[1878] := 0.1851012;
   Prof_PriceDA.Data[1879] := 0.1851012;
   Prof_PriceDA.Data[1880] := 0.2071332;
   Prof_PriceDA.Data[1881] := 0.2071332;
   Prof_PriceDA.Data[1882] := 0.2071332;
   Prof_PriceDA.Data[1883] := 0.2071332;
   Prof_PriceDA.Data[1884] := 0.2981016;
   Prof_PriceDA.Data[1885] := 0.2981016;
   Prof_PriceDA.Data[1886] := 0.2981016;
   Prof_PriceDA.Data[1887] := 0.2981016;
   Prof_PriceDA.Data[1888] := 0.446472;
   Prof_PriceDA.Data[1889] := 0.446472;
   Prof_PriceDA.Data[1890] := 0.446472;
   Prof_PriceDA.Data[1891] := 0.446472;
   Prof_PriceDA.Data[1892] := 0.6208812;
   Prof_PriceDA.Data[1893] := 0.6208812;
   Prof_PriceDA.Data[1894] := 0.6208812;
   Prof_PriceDA.Data[1895] := 0.6208812;
   Prof_PriceDA.Data[1896] := 0.5111424;
   Prof_PriceDA.Data[1897] := 0.5111424;
   Prof_PriceDA.Data[1898] := 0.5111424;
   Prof_PriceDA.Data[1899] := 0.5111424;
   Prof_PriceDA.Data[1900] := 0.3192156;
   Prof_PriceDA.Data[1901] := 0.3192156;
   Prof_PriceDA.Data[1902] := 0.3192156;
   Prof_PriceDA.Data[1903] := 0.3192156;
   Prof_PriceDA.Data[1904] := 0.2376;
   Prof_PriceDA.Data[1905] := 0.2376;
   Prof_PriceDA.Data[1906] := 0.2376;
   Prof_PriceDA.Data[1907] := 0.2376;
   Prof_PriceDA.Data[1908] := 0.1836;
   Prof_PriceDA.Data[1909] := 0.1836;
   Prof_PriceDA.Data[1910] := 0.1836;
   Prof_PriceDA.Data[1911] := 0.1836;
   Prof_PriceDA.Data[1912] := 0.1718928;
   Prof_PriceDA.Data[1913] := 0.1718928;
   Prof_PriceDA.Data[1914] := 0.1718928;
   Prof_PriceDA.Data[1915] := 0.1718928;
   Prof_PriceDA.Data[1916] := 0.1540944;
   Prof_PriceDA.Data[1917] := 0.1540944;
   Prof_PriceDA.Data[1918] := 0.1540944;
   Prof_PriceDA.Data[1919] := 0.1540944;
   Prof_PriceDA.Data[1920] := 0.1477764;
   Prof_PriceDA.Data[1921] := 0.1477764;
   Prof_PriceDA.Data[1922] := 0.1477764;
   Prof_PriceDA.Data[1923] := 0.1477764;
   Prof_PriceDA.Data[1924] := 0.1417932;
   Prof_PriceDA.Data[1925] := 0.1417932;
   Prof_PriceDA.Data[1926] := 0.1417932;
   Prof_PriceDA.Data[1927] := 0.1417932;
   Prof_PriceDA.Data[1928] := 0.134622;
   Prof_PriceDA.Data[1929] := 0.134622;
   Prof_PriceDA.Data[1930] := 0.134622;
   Prof_PriceDA.Data[1931] := 0.134622;
   Prof_PriceDA.Data[1932] := 0.1350972;
   Prof_PriceDA.Data[1933] := 0.1350972;
   Prof_PriceDA.Data[1934] := 0.1350972;
   Prof_PriceDA.Data[1935] := 0.1350972;
   Prof_PriceDA.Data[1936] := 0.1429056;
   Prof_PriceDA.Data[1937] := 0.1429056;
   Prof_PriceDA.Data[1938] := 0.1429056;
   Prof_PriceDA.Data[1939] := 0.1429056;
   Prof_PriceDA.Data[1940] := 0.16416;
   Prof_PriceDA.Data[1941] := 0.16416;
   Prof_PriceDA.Data[1942] := 0.16416;
   Prof_PriceDA.Data[1943] := 0.16416;
   Prof_PriceDA.Data[1944] := 0.207414;
   Prof_PriceDA.Data[1945] := 0.207414;
   Prof_PriceDA.Data[1946] := 0.207414;
   Prof_PriceDA.Data[1947] := 0.207414;
   Prof_PriceDA.Data[1948] := 0.3141612;
   Prof_PriceDA.Data[1949] := 0.3141612;
   Prof_PriceDA.Data[1950] := 0.3141612;
   Prof_PriceDA.Data[1951] := 0.3141612;
   Prof_PriceDA.Data[1952] := 0.4177224;
   Prof_PriceDA.Data[1953] := 0.4177224;
   Prof_PriceDA.Data[1954] := 0.4177224;
   Prof_PriceDA.Data[1955] := 0.4177224;
   Prof_PriceDA.Data[1956] := 0.2861676;
   Prof_PriceDA.Data[1957] := 0.2861676;
   Prof_PriceDA.Data[1958] := 0.2861676;
   Prof_PriceDA.Data[1959] := 0.2861676;
   Prof_PriceDA.Data[1960] := 0.2540484;
   Prof_PriceDA.Data[1961] := 0.2540484;
   Prof_PriceDA.Data[1962] := 0.2540484;
   Prof_PriceDA.Data[1963] := 0.2540484;
   Prof_PriceDA.Data[1964] := 0.2179224;
   Prof_PriceDA.Data[1965] := 0.2179224;
   Prof_PriceDA.Data[1966] := 0.2179224;
   Prof_PriceDA.Data[1967] := 0.2179224;
   Prof_PriceDA.Data[1968] := 0.2129004;
   Prof_PriceDA.Data[1969] := 0.2129004;
   Prof_PriceDA.Data[1970] := 0.2129004;
   Prof_PriceDA.Data[1971] := 0.2129004;
   Prof_PriceDA.Data[1972] := 0.1951344;
   Prof_PriceDA.Data[1973] := 0.1951344;
   Prof_PriceDA.Data[1974] := 0.1951344;
   Prof_PriceDA.Data[1975] := 0.1951344;
   Prof_PriceDA.Data[1976] := 0.2188512;
   Prof_PriceDA.Data[1977] := 0.2188512;
   Prof_PriceDA.Data[1978] := 0.2188512;
   Prof_PriceDA.Data[1979] := 0.2188512;
   Prof_PriceDA.Data[1980] := 0.3057588;
   Prof_PriceDA.Data[1981] := 0.3057588;
   Prof_PriceDA.Data[1982] := 0.3057588;
   Prof_PriceDA.Data[1983] := 0.3057588;
   Prof_PriceDA.Data[1984] := 0.245214;
   Prof_PriceDA.Data[1985] := 0.245214;
   Prof_PriceDA.Data[1986] := 0.245214;
   Prof_PriceDA.Data[1987] := 0.245214;
   Prof_PriceDA.Data[1988] := 0.3387744;
   Prof_PriceDA.Data[1989] := 0.3387744;
   Prof_PriceDA.Data[1990] := 0.3387744;
   Prof_PriceDA.Data[1991] := 0.3387744;
   Prof_PriceDA.Data[1992] := 0.2779704;
   Prof_PriceDA.Data[1993] := 0.2779704;
   Prof_PriceDA.Data[1994] := 0.2779704;
   Prof_PriceDA.Data[1995] := 0.2779704;
   Prof_PriceDA.Data[1996] := 0.2207844;
   Prof_PriceDA.Data[1997] := 0.2207844;
   Prof_PriceDA.Data[1998] := 0.2207844;
   Prof_PriceDA.Data[1999] := 0.2207844;
   Prof_PriceDA.Data[2000] := 0.190728;
   Prof_PriceDA.Data[2001] := 0.190728;
   Prof_PriceDA.Data[2002] := 0.190728;
   Prof_PriceDA.Data[2003] := 0.190728;
   Prof_PriceDA.Data[2004] := 0.1687392;
   Prof_PriceDA.Data[2005] := 0.1687392;
   Prof_PriceDA.Data[2006] := 0.1687392;
   Prof_PriceDA.Data[2007] := 0.1687392;
   Prof_PriceDA.Data[2008] := 0.153684;
   Prof_PriceDA.Data[2009] := 0.153684;
   Prof_PriceDA.Data[2010] := 0.153684;
   Prof_PriceDA.Data[2011] := 0.153684;
   Prof_PriceDA.Data[2012] := 0.144234;
   Prof_PriceDA.Data[2013] := 0.144234;
   Prof_PriceDA.Data[2014] := 0.144234;
   Prof_PriceDA.Data[2015] := 0.144234;
   Prof_PriceDA.Data[2016] := 0.141588;
   Prof_PriceDA.Data[2017] := 0.141588;
   Prof_PriceDA.Data[2018] := 0.141588;
   Prof_PriceDA.Data[2019] := 0.141588;
   Prof_PriceDA.Data[2020] := 0.1360152;
   Prof_PriceDA.Data[2021] := 0.1360152;
   Prof_PriceDA.Data[2022] := 0.1360152;
   Prof_PriceDA.Data[2023] := 0.1360152;
   Prof_PriceDA.Data[2024] := 0.1345896;
   Prof_PriceDA.Data[2025] := 0.1345896;
   Prof_PriceDA.Data[2026] := 0.1345896;
   Prof_PriceDA.Data[2027] := 0.1345896;
   Prof_PriceDA.Data[2028] := 0.1350972;
   Prof_PriceDA.Data[2029] := 0.1350972;
   Prof_PriceDA.Data[2030] := 0.1350972;
   Prof_PriceDA.Data[2031] := 0.1350972;
   Prof_PriceDA.Data[2032] := 0.1372464;
   Prof_PriceDA.Data[2033] := 0.1372464;
   Prof_PriceDA.Data[2034] := 0.1372464;
   Prof_PriceDA.Data[2035] := 0.1372464;
   Prof_PriceDA.Data[2036] := 0.1506816;
   Prof_PriceDA.Data[2037] := 0.1506816;
   Prof_PriceDA.Data[2038] := 0.1506816;
   Prof_PriceDA.Data[2039] := 0.1506816;
   Prof_PriceDA.Data[2040] := 0.20925;
   Prof_PriceDA.Data[2041] := 0.20925;
   Prof_PriceDA.Data[2042] := 0.20925;
   Prof_PriceDA.Data[2043] := 0.20925;
   Prof_PriceDA.Data[2044] := 0.3410964;
   Prof_PriceDA.Data[2045] := 0.3410964;
   Prof_PriceDA.Data[2046] := 0.3410964;
   Prof_PriceDA.Data[2047] := 0.3410964;
   Prof_PriceDA.Data[2048] := 0.2672136;
   Prof_PriceDA.Data[2049] := 0.2672136;
   Prof_PriceDA.Data[2050] := 0.2672136;
   Prof_PriceDA.Data[2051] := 0.2672136;
   Prof_PriceDA.Data[2052] := 0.2153628;
   Prof_PriceDA.Data[2053] := 0.2153628;
   Prof_PriceDA.Data[2054] := 0.2153628;
   Prof_PriceDA.Data[2055] := 0.2153628;
   Prof_PriceDA.Data[2056] := 0.1933848;
   Prof_PriceDA.Data[2057] := 0.1933848;
   Prof_PriceDA.Data[2058] := 0.1933848;
   Prof_PriceDA.Data[2059] := 0.1933848;
   Prof_PriceDA.Data[2060] := 0.1867752;
   Prof_PriceDA.Data[2061] := 0.1867752;
   Prof_PriceDA.Data[2062] := 0.1867752;
   Prof_PriceDA.Data[2063] := 0.1867752;
   Prof_PriceDA.Data[2064] := 0.1782;
   Prof_PriceDA.Data[2065] := 0.1782;
   Prof_PriceDA.Data[2066] := 0.1782;
   Prof_PriceDA.Data[2067] := 0.1782;
   Prof_PriceDA.Data[2068] := 0.1836;
   Prof_PriceDA.Data[2069] := 0.1836;
   Prof_PriceDA.Data[2070] := 0.1836;
   Prof_PriceDA.Data[2071] := 0.1836;
   Prof_PriceDA.Data[2072] := 0.1943136;
   Prof_PriceDA.Data[2073] := 0.1943136;
   Prof_PriceDA.Data[2074] := 0.1943136;
   Prof_PriceDA.Data[2075] := 0.1943136;
   Prof_PriceDA.Data[2076] := 0.2137752;
   Prof_PriceDA.Data[2077] := 0.2137752;
   Prof_PriceDA.Data[2078] := 0.2137752;
   Prof_PriceDA.Data[2079] := 0.2137752;
   Prof_PriceDA.Data[2080] := 0.2703888;
   Prof_PriceDA.Data[2081] := 0.2703888;
   Prof_PriceDA.Data[2082] := 0.2703888;
   Prof_PriceDA.Data[2083] := 0.2703888;
   Prof_PriceDA.Data[2084] := 0.276102;
   Prof_PriceDA.Data[2085] := 0.276102;
   Prof_PriceDA.Data[2086] := 0.276102;
   Prof_PriceDA.Data[2087] := 0.276102;
   Prof_PriceDA.Data[2088] := 0.2261952;
   Prof_PriceDA.Data[2089] := 0.2261952;
   Prof_PriceDA.Data[2090] := 0.2261952;
   Prof_PriceDA.Data[2091] := 0.2261952;
   Prof_PriceDA.Data[2092] := 0.222642;
   Prof_PriceDA.Data[2093] := 0.222642;
   Prof_PriceDA.Data[2094] := 0.222642;
   Prof_PriceDA.Data[2095] := 0.222642;
   Prof_PriceDA.Data[2096] := 0.2220156;
   Prof_PriceDA.Data[2097] := 0.2220156;
   Prof_PriceDA.Data[2098] := 0.2220156;
   Prof_PriceDA.Data[2099] := 0.2220156;
   Prof_PriceDA.Data[2100] := 0.1710072;
   Prof_PriceDA.Data[2101] := 0.1710072;
   Prof_PriceDA.Data[2102] := 0.1710072;
   Prof_PriceDA.Data[2103] := 0.1710072;
   Prof_PriceDA.Data[2104] := 0.1589436;
   Prof_PriceDA.Data[2105] := 0.1589436;
   Prof_PriceDA.Data[2106] := 0.1589436;
   Prof_PriceDA.Data[2107] := 0.1589436;
   Prof_PriceDA.Data[2108] := 0.145854;
   Prof_PriceDA.Data[2109] := 0.145854;
   Prof_PriceDA.Data[2110] := 0.145854;
   Prof_PriceDA.Data[2111] := 0.145854;
   Prof_PriceDA.Data[2112] := 0.1353888;
   Prof_PriceDA.Data[2113] := 0.1353888;
   Prof_PriceDA.Data[2114] := 0.1353888;
   Prof_PriceDA.Data[2115] := 0.1353888;
   Prof_PriceDA.Data[2116] := 0.1299564;
   Prof_PriceDA.Data[2117] := 0.1299564;
   Prof_PriceDA.Data[2118] := 0.1299564;
   Prof_PriceDA.Data[2119] := 0.1299564;
   Prof_PriceDA.Data[2120] := 0.119394;
   Prof_PriceDA.Data[2121] := 0.119394;
   Prof_PriceDA.Data[2122] := 0.119394;
   Prof_PriceDA.Data[2123] := 0.119394;
   Prof_PriceDA.Data[2124] := 0.1175796;
   Prof_PriceDA.Data[2125] := 0.1175796;
   Prof_PriceDA.Data[2126] := 0.1175796;
   Prof_PriceDA.Data[2127] := 0.1175796;
   Prof_PriceDA.Data[2128] := 0.1227096;
   Prof_PriceDA.Data[2129] := 0.1227096;
   Prof_PriceDA.Data[2130] := 0.1227096;
   Prof_PriceDA.Data[2131] := 0.1227096;
   Prof_PriceDA.Data[2132] := 0.1344708;
   Prof_PriceDA.Data[2133] := 0.1344708;
   Prof_PriceDA.Data[2134] := 0.1344708;
   Prof_PriceDA.Data[2135] := 0.1344708;
   Prof_PriceDA.Data[2136] := 0.1809864;
   Prof_PriceDA.Data[2137] := 0.1809864;
   Prof_PriceDA.Data[2138] := 0.1809864;
   Prof_PriceDA.Data[2139] := 0.1809864;
   Prof_PriceDA.Data[2140] := 0.2092608;
   Prof_PriceDA.Data[2141] := 0.2092608;
   Prof_PriceDA.Data[2142] := 0.2092608;
   Prof_PriceDA.Data[2143] := 0.2092608;
   Prof_PriceDA.Data[2144] := 0.1881684;
   Prof_PriceDA.Data[2145] := 0.1881684;
   Prof_PriceDA.Data[2146] := 0.1881684;
   Prof_PriceDA.Data[2147] := 0.1881684;
   Prof_PriceDA.Data[2148] := 0.1808568;
   Prof_PriceDA.Data[2149] := 0.1808568;
   Prof_PriceDA.Data[2150] := 0.1808568;
   Prof_PriceDA.Data[2151] := 0.1808568;
   Prof_PriceDA.Data[2152] := 0.1625292;
   Prof_PriceDA.Data[2153] := 0.1625292;
   Prof_PriceDA.Data[2154] := 0.1625292;
   Prof_PriceDA.Data[2155] := 0.1625292;
   Prof_PriceDA.Data[2156] := 0.1594728;
   Prof_PriceDA.Data[2157] := 0.1594728;
   Prof_PriceDA.Data[2158] := 0.1594728;
   Prof_PriceDA.Data[2159] := 0.1594728;
   Prof_PriceDA.Data[2160] := 0.1543104;
   Prof_PriceDA.Data[2161] := 0.1543104;
   Prof_PriceDA.Data[2162] := 0.1543104;
   Prof_PriceDA.Data[2163] := 0.1543104;
   Prof_PriceDA.Data[2164] := 0.1588032;
   Prof_PriceDA.Data[2165] := 0.1588032;
   Prof_PriceDA.Data[2166] := 0.1588032;
   Prof_PriceDA.Data[2167] := 0.1588032;
   Prof_PriceDA.Data[2168] := 0.1690416;
   Prof_PriceDA.Data[2169] := 0.1690416;
   Prof_PriceDA.Data[2170] := 0.1690416;
   Prof_PriceDA.Data[2171] := 0.1690416;
   Prof_PriceDA.Data[2172] := 0.1919376;
   Prof_PriceDA.Data[2173] := 0.1919376;
   Prof_PriceDA.Data[2174] := 0.1919376;
   Prof_PriceDA.Data[2175] := 0.1919376;
   Prof_PriceDA.Data[2176] := 0.2108916;
   Prof_PriceDA.Data[2177] := 0.2108916;
   Prof_PriceDA.Data[2178] := 0.2108916;
   Prof_PriceDA.Data[2179] := 0.2108916;
   Prof_PriceDA.Data[2180] := 0.2148012;
   Prof_PriceDA.Data[2181] := 0.2148012;
   Prof_PriceDA.Data[2182] := 0.2148012;
   Prof_PriceDA.Data[2183] := 0.2148012;
   Prof_PriceDA.Data[2184] := 0.2028672;
   Prof_PriceDA.Data[2185] := 0.2028672;
   Prof_PriceDA.Data[2186] := 0.2028672;
   Prof_PriceDA.Data[2187] := 0.2028672;
   Prof_PriceDA.Data[2188] := 0.1957824;
   Prof_PriceDA.Data[2189] := 0.1957824;
   Prof_PriceDA.Data[2190] := 0.1957824;
   Prof_PriceDA.Data[2191] := 0.1957824;
   Prof_PriceDA.Data[2192] := 0.2018628;
   Prof_PriceDA.Data[2193] := 0.2018628;
   Prof_PriceDA.Data[2194] := 0.2018628;
   Prof_PriceDA.Data[2195] := 0.2018628;
   Prof_PriceDA.Data[2196] := 0.1633608;
   Prof_PriceDA.Data[2197] := 0.1633608;
   Prof_PriceDA.Data[2198] := 0.1633608;
   Prof_PriceDA.Data[2199] := 0.1633608;
   Prof_PriceDA.Data[2200] := 0.1606176;
   Prof_PriceDA.Data[2201] := 0.1606176;
   Prof_PriceDA.Data[2202] := 0.1606176;
   Prof_PriceDA.Data[2203] := 0.1606176;
   Prof_PriceDA.Data[2204] := 0.136188;
   Prof_PriceDA.Data[2205] := 0.136188;
   Prof_PriceDA.Data[2206] := 0.136188;
   Prof_PriceDA.Data[2207] := 0.136188;
   Prof_PriceDA.Data[2208] := 0.127656;
   Prof_PriceDA.Data[2209] := 0.127656;
   Prof_PriceDA.Data[2210] := 0.127656;
   Prof_PriceDA.Data[2211] := 0.127656;
   Prof_PriceDA.Data[2212] := 0.1162512;
   Prof_PriceDA.Data[2213] := 0.1162512;
   Prof_PriceDA.Data[2214] := 0.1162512;
   Prof_PriceDA.Data[2215] := 0.1162512;
   Prof_PriceDA.Data[2216] := 0.1107;
   Prof_PriceDA.Data[2217] := 0.1107;
   Prof_PriceDA.Data[2218] := 0.1107;
   Prof_PriceDA.Data[2219] := 0.1107;
   Prof_PriceDA.Data[2220] := 0.1093392;
   Prof_PriceDA.Data[2221] := 0.1093392;
   Prof_PriceDA.Data[2222] := 0.1093392;
   Prof_PriceDA.Data[2223] := 0.1093392;
   Prof_PriceDA.Data[2224] := 0.1170288;
   Prof_PriceDA.Data[2225] := 0.1170288;
   Prof_PriceDA.Data[2226] := 0.1170288;
   Prof_PriceDA.Data[2227] := 0.1170288;
   Prof_PriceDA.Data[2228] := 0.1424304;
   Prof_PriceDA.Data[2229] := 0.1424304;
   Prof_PriceDA.Data[2230] := 0.1424304;
   Prof_PriceDA.Data[2231] := 0.1424304;
   Prof_PriceDA.Data[2232] := 0.17469;
   Prof_PriceDA.Data[2233] := 0.17469;
   Prof_PriceDA.Data[2234] := 0.17469;
   Prof_PriceDA.Data[2235] := 0.17469;
   Prof_PriceDA.Data[2236] := 0.1909872;
   Prof_PriceDA.Data[2237] := 0.1909872;
   Prof_PriceDA.Data[2238] := 0.1909872;
   Prof_PriceDA.Data[2239] := 0.1909872;
   Prof_PriceDA.Data[2240] := 0.1764828;
   Prof_PriceDA.Data[2241] := 0.1764828;
   Prof_PriceDA.Data[2242] := 0.1764828;
   Prof_PriceDA.Data[2243] := 0.1764828;
   Prof_PriceDA.Data[2244] := 0.1599048;
   Prof_PriceDA.Data[2245] := 0.1599048;
   Prof_PriceDA.Data[2246] := 0.1599048;
   Prof_PriceDA.Data[2247] := 0.1599048;
   Prof_PriceDA.Data[2248] := 0.1535652;
   Prof_PriceDA.Data[2249] := 0.1535652;
   Prof_PriceDA.Data[2250] := 0.1535652;
   Prof_PriceDA.Data[2251] := 0.1535652;
   Prof_PriceDA.Data[2252] := 0.1422576;
   Prof_PriceDA.Data[2253] := 0.1422576;
   Prof_PriceDA.Data[2254] := 0.1422576;
   Prof_PriceDA.Data[2255] := 0.1422576;
   Prof_PriceDA.Data[2256] := 0.1392444;
   Prof_PriceDA.Data[2257] := 0.1392444;
   Prof_PriceDA.Data[2258] := 0.1392444;
   Prof_PriceDA.Data[2259] := 0.1392444;
   Prof_PriceDA.Data[2260] := 0.13662;
   Prof_PriceDA.Data[2261] := 0.13662;
   Prof_PriceDA.Data[2262] := 0.13662;
   Prof_PriceDA.Data[2263] := 0.13662;
   Prof_PriceDA.Data[2264] := 0.1417716;
   Prof_PriceDA.Data[2265] := 0.1417716;
   Prof_PriceDA.Data[2266] := 0.1417716;
   Prof_PriceDA.Data[2267] := 0.1417716;
   Prof_PriceDA.Data[2268] := 0.161892;
   Prof_PriceDA.Data[2269] := 0.161892;
   Prof_PriceDA.Data[2270] := 0.161892;
   Prof_PriceDA.Data[2271] := 0.161892;
   Prof_PriceDA.Data[2272] := 0.1961064;
   Prof_PriceDA.Data[2273] := 0.1961064;
   Prof_PriceDA.Data[2274] := 0.1961064;
   Prof_PriceDA.Data[2275] := 0.1961064;
   Prof_PriceDA.Data[2276] := 0.1983744;
   Prof_PriceDA.Data[2277] := 0.1983744;
   Prof_PriceDA.Data[2278] := 0.1983744;
   Prof_PriceDA.Data[2279] := 0.1983744;
   Prof_PriceDA.Data[2280] := 0.1922616;
   Prof_PriceDA.Data[2281] := 0.1922616;
   Prof_PriceDA.Data[2282] := 0.1922616;
   Prof_PriceDA.Data[2283] := 0.1922616;
   Prof_PriceDA.Data[2284] := 0.1883412;
   Prof_PriceDA.Data[2285] := 0.1883412;
   Prof_PriceDA.Data[2286] := 0.1883412;
   Prof_PriceDA.Data[2287] := 0.1883412;
   Prof_PriceDA.Data[2288] := 0.1774872;
   Prof_PriceDA.Data[2289] := 0.1774872;
   Prof_PriceDA.Data[2290] := 0.1774872;
   Prof_PriceDA.Data[2291] := 0.1774872;
   Prof_PriceDA.Data[2292] := 0.1666008;
   Prof_PriceDA.Data[2293] := 0.1666008;
   Prof_PriceDA.Data[2294] := 0.1666008;
   Prof_PriceDA.Data[2295] := 0.1666008;
   Prof_PriceDA.Data[2296] := 0.1547208;
   Prof_PriceDA.Data[2297] := 0.1547208;
   Prof_PriceDA.Data[2298] := 0.1547208;
   Prof_PriceDA.Data[2299] := 0.1547208;
   Prof_PriceDA.Data[2300] := 0.1429488;
   Prof_PriceDA.Data[2301] := 0.1429488;
   Prof_PriceDA.Data[2302] := 0.1429488;
   Prof_PriceDA.Data[2303] := 0.1429488;
   Prof_PriceDA.Data[2304] := 0.1203336;
   Prof_PriceDA.Data[2305] := 0.1203336;
   Prof_PriceDA.Data[2306] := 0.1203336;
   Prof_PriceDA.Data[2307] := 0.1203336;
   Prof_PriceDA.Data[2308] := 0.1117476;
   Prof_PriceDA.Data[2309] := 0.1117476;
   Prof_PriceDA.Data[2310] := 0.1117476;
   Prof_PriceDA.Data[2311] := 0.1117476;
   Prof_PriceDA.Data[2312] := 0.0980856;
   Prof_PriceDA.Data[2313] := 0.0980856;
   Prof_PriceDA.Data[2314] := 0.0980856;
   Prof_PriceDA.Data[2315] := 0.0980856;
   Prof_PriceDA.Data[2316] := 0.094878;
   Prof_PriceDA.Data[2317] := 0.094878;
   Prof_PriceDA.Data[2318] := 0.094878;
   Prof_PriceDA.Data[2319] := 0.094878;
   Prof_PriceDA.Data[2320] := 0.0971136;
   Prof_PriceDA.Data[2321] := 0.0971136;
   Prof_PriceDA.Data[2322] := 0.0971136;
   Prof_PriceDA.Data[2323] := 0.0971136;
   Prof_PriceDA.Data[2324] := 0.1055808;
   Prof_PriceDA.Data[2325] := 0.1055808;
   Prof_PriceDA.Data[2326] := 0.1055808;
   Prof_PriceDA.Data[2327] := 0.1055808;
   Prof_PriceDA.Data[2328] := 0.1218564;
   Prof_PriceDA.Data[2329] := 0.1218564;
   Prof_PriceDA.Data[2330] := 0.1218564;
   Prof_PriceDA.Data[2331] := 0.1218564;
   Prof_PriceDA.Data[2332] := 0.1337904;
   Prof_PriceDA.Data[2333] := 0.1337904;
   Prof_PriceDA.Data[2334] := 0.1337904;
   Prof_PriceDA.Data[2335] := 0.1337904;
   Prof_PriceDA.Data[2336] := 0.1181628;
   Prof_PriceDA.Data[2337] := 0.1181628;
   Prof_PriceDA.Data[2338] := 0.1181628;
   Prof_PriceDA.Data[2339] := 0.1181628;
   Prof_PriceDA.Data[2340] := 0.1153224;
   Prof_PriceDA.Data[2341] := 0.1153224;
   Prof_PriceDA.Data[2342] := 0.1153224;
   Prof_PriceDA.Data[2343] := 0.1153224;
   Prof_PriceDA.Data[2344] := 0.1033776;
   Prof_PriceDA.Data[2345] := 0.1033776;
   Prof_PriceDA.Data[2346] := 0.1033776;
   Prof_PriceDA.Data[2347] := 0.1033776;
   Prof_PriceDA.Data[2348] := 0.0975888;
   Prof_PriceDA.Data[2349] := 0.0975888;
   Prof_PriceDA.Data[2350] := 0.0975888;
   Prof_PriceDA.Data[2351] := 0.0975888;
   Prof_PriceDA.Data[2352] := 0.09396;
   Prof_PriceDA.Data[2353] := 0.09396;
   Prof_PriceDA.Data[2354] := 0.09396;
   Prof_PriceDA.Data[2355] := 0.09396;
   Prof_PriceDA.Data[2356] := 0.0924372;
   Prof_PriceDA.Data[2357] := 0.0924372;
   Prof_PriceDA.Data[2358] := 0.0924372;
   Prof_PriceDA.Data[2359] := 0.0924372;
   Prof_PriceDA.Data[2360] := 0.1067256;
   Prof_PriceDA.Data[2361] := 0.1067256;
   Prof_PriceDA.Data[2362] := 0.1067256;
   Prof_PriceDA.Data[2363] := 0.1067256;
   Prof_PriceDA.Data[2364] := 0.1288872;
   Prof_PriceDA.Data[2365] := 0.1288872;
   Prof_PriceDA.Data[2366] := 0.1288872;
   Prof_PriceDA.Data[2367] := 0.1288872;
   Prof_PriceDA.Data[2368] := 0.1661148;
   Prof_PriceDA.Data[2369] := 0.1661148;
   Prof_PriceDA.Data[2370] := 0.1661148;
   Prof_PriceDA.Data[2371] := 0.1661148;
   Prof_PriceDA.Data[2372] := 0.1701108;
   Prof_PriceDA.Data[2373] := 0.1701108;
   Prof_PriceDA.Data[2374] := 0.1701108;
   Prof_PriceDA.Data[2375] := 0.1701108;
   Prof_PriceDA.Data[2376] := 0.1716444;
   Prof_PriceDA.Data[2377] := 0.1716444;
   Prof_PriceDA.Data[2378] := 0.1716444;
   Prof_PriceDA.Data[2379] := 0.1716444;
   Prof_PriceDA.Data[2380] := 0.1709208;
   Prof_PriceDA.Data[2381] := 0.1709208;
   Prof_PriceDA.Data[2382] := 0.1709208;
   Prof_PriceDA.Data[2383] := 0.1709208;
   Prof_PriceDA.Data[2384] := 0.162864;
   Prof_PriceDA.Data[2385] := 0.162864;
   Prof_PriceDA.Data[2386] := 0.162864;
   Prof_PriceDA.Data[2387] := 0.162864;
   Prof_PriceDA.Data[2388] := 0.155574;
   Prof_PriceDA.Data[2389] := 0.155574;
   Prof_PriceDA.Data[2390] := 0.155574;
   Prof_PriceDA.Data[2391] := 0.155574;
   Prof_PriceDA.Data[2392] := 0.1481004;
   Prof_PriceDA.Data[2393] := 0.1481004;
   Prof_PriceDA.Data[2394] := 0.1481004;
   Prof_PriceDA.Data[2395] := 0.1481004;
   Prof_PriceDA.Data[2396] := 0.135;
   Prof_PriceDA.Data[2397] := 0.135;
   Prof_PriceDA.Data[2398] := 0.135;
   Prof_PriceDA.Data[2399] := 0.135;
   Prof_PriceDA.Data[2400] := 0.1419552;
   Prof_PriceDA.Data[2401] := 0.1419552;
   Prof_PriceDA.Data[2402] := 0.1419552;
   Prof_PriceDA.Data[2403] := 0.1419552;
   Prof_PriceDA.Data[2404] := 0.1297404;
   Prof_PriceDA.Data[2405] := 0.1297404;
   Prof_PriceDA.Data[2406] := 0.1297404;
   Prof_PriceDA.Data[2407] := 0.1297404;
   Prof_PriceDA.Data[2408] := 0.1272888;
   Prof_PriceDA.Data[2409] := 0.1272888;
   Prof_PriceDA.Data[2410] := 0.1272888;
   Prof_PriceDA.Data[2411] := 0.1272888;
   Prof_PriceDA.Data[2412] := 0.1204524;
   Prof_PriceDA.Data[2413] := 0.1204524;
   Prof_PriceDA.Data[2414] := 0.1204524;
   Prof_PriceDA.Data[2415] := 0.1204524;
   Prof_PriceDA.Data[2416] := 0.12096;
   Prof_PriceDA.Data[2417] := 0.12096;
   Prof_PriceDA.Data[2418] := 0.12096;
   Prof_PriceDA.Data[2419] := 0.12096;
   Prof_PriceDA.Data[2420] := 0.1231524;
   Prof_PriceDA.Data[2421] := 0.1231524;
   Prof_PriceDA.Data[2422] := 0.1231524;
   Prof_PriceDA.Data[2423] := 0.1231524;
   Prof_PriceDA.Data[2424] := 0.1255176;
   Prof_PriceDA.Data[2425] := 0.1255176;
   Prof_PriceDA.Data[2426] := 0.1255176;
   Prof_PriceDA.Data[2427] := 0.1255176;
   Prof_PriceDA.Data[2428] := 0.1334664;
   Prof_PriceDA.Data[2429] := 0.1334664;
   Prof_PriceDA.Data[2430] := 0.1334664;
   Prof_PriceDA.Data[2431] := 0.1334664;
   Prof_PriceDA.Data[2432] := 0.1427112;
   Prof_PriceDA.Data[2433] := 0.1427112;
   Prof_PriceDA.Data[2434] := 0.1427112;
   Prof_PriceDA.Data[2435] := 0.1427112;
   Prof_PriceDA.Data[2436] := 0.1400004;
   Prof_PriceDA.Data[2437] := 0.1400004;
   Prof_PriceDA.Data[2438] := 0.1400004;
   Prof_PriceDA.Data[2439] := 0.1400004;
   Prof_PriceDA.Data[2440] := 0.1207656;
   Prof_PriceDA.Data[2441] := 0.1207656;
   Prof_PriceDA.Data[2442] := 0.1207656;
   Prof_PriceDA.Data[2443] := 0.1207656;
   Prof_PriceDA.Data[2444] := 0.112752;
   Prof_PriceDA.Data[2445] := 0.112752;
   Prof_PriceDA.Data[2446] := 0.112752;
   Prof_PriceDA.Data[2447] := 0.112752;
   Prof_PriceDA.Data[2448] := 0.1054188;
   Prof_PriceDA.Data[2449] := 0.1054188;
   Prof_PriceDA.Data[2450] := 0.1054188;
   Prof_PriceDA.Data[2451] := 0.1054188;
   Prof_PriceDA.Data[2452] := 0.1028808;
   Prof_PriceDA.Data[2453] := 0.1028808;
   Prof_PriceDA.Data[2454] := 0.1028808;
   Prof_PriceDA.Data[2455] := 0.1028808;
   Prof_PriceDA.Data[2456] := 0.1209168;
   Prof_PriceDA.Data[2457] := 0.1209168;
   Prof_PriceDA.Data[2458] := 0.1209168;
   Prof_PriceDA.Data[2459] := 0.1209168;
   Prof_PriceDA.Data[2460] := 0.13095;
   Prof_PriceDA.Data[2461] := 0.13095;
   Prof_PriceDA.Data[2462] := 0.13095;
   Prof_PriceDA.Data[2463] := 0.13095;
   Prof_PriceDA.Data[2464] := 0.1467288;
   Prof_PriceDA.Data[2465] := 0.1467288;
   Prof_PriceDA.Data[2466] := 0.1467288;
   Prof_PriceDA.Data[2467] := 0.1467288;
   Prof_PriceDA.Data[2468] := 0.1559088;
   Prof_PriceDA.Data[2469] := 0.1559088;
   Prof_PriceDA.Data[2470] := 0.1559088;
   Prof_PriceDA.Data[2471] := 0.1559088;
   Prof_PriceDA.Data[2472] := 0.1424628;
   Prof_PriceDA.Data[2473] := 0.1424628;
   Prof_PriceDA.Data[2474] := 0.1424628;
   Prof_PriceDA.Data[2475] := 0.1424628;
   Prof_PriceDA.Data[2476] := 0.1443312;
   Prof_PriceDA.Data[2477] := 0.1443312;
   Prof_PriceDA.Data[2478] := 0.1443312;
   Prof_PriceDA.Data[2479] := 0.1443312;
   Prof_PriceDA.Data[2480] := 0.1348812;
   Prof_PriceDA.Data[2481] := 0.1348812;
   Prof_PriceDA.Data[2482] := 0.1348812;
   Prof_PriceDA.Data[2483] := 0.1348812;
   Prof_PriceDA.Data[2484] := 0.1245888;
   Prof_PriceDA.Data[2485] := 0.1245888;
   Prof_PriceDA.Data[2486] := 0.1245888;
   Prof_PriceDA.Data[2487] := 0.1245888;
   Prof_PriceDA.Data[2488] := 0.104004;
   Prof_PriceDA.Data[2489] := 0.104004;
   Prof_PriceDA.Data[2490] := 0.104004;
   Prof_PriceDA.Data[2491] := 0.104004;
   Prof_PriceDA.Data[2492] := 0.08397;
   Prof_PriceDA.Data[2493] := 0.08397;
   Prof_PriceDA.Data[2494] := 0.08397;
   Prof_PriceDA.Data[2495] := 0.08397;
   Prof_PriceDA.Data[2496] := 0.0654696;
   Prof_PriceDA.Data[2497] := 0.0654696;
   Prof_PriceDA.Data[2498] := 0.0654696;
   Prof_PriceDA.Data[2499] := 0.0654696;
   Prof_PriceDA.Data[2500] := 0.0605124;
   Prof_PriceDA.Data[2501] := 0.0605124;
   Prof_PriceDA.Data[2502] := 0.0605124;
   Prof_PriceDA.Data[2503] := 0.0605124;
   Prof_PriceDA.Data[2504] := 0.0433404;
   Prof_PriceDA.Data[2505] := 0.0433404;
   Prof_PriceDA.Data[2506] := 0.0433404;
   Prof_PriceDA.Data[2507] := 0.0433404;
   Prof_PriceDA.Data[2508] := 0.032022;
   Prof_PriceDA.Data[2509] := 0.032022;
   Prof_PriceDA.Data[2510] := 0.032022;
   Prof_PriceDA.Data[2511] := 0.032022;
   Prof_PriceDA.Data[2512] := 0.0490536;
   Prof_PriceDA.Data[2513] := 0.0490536;
   Prof_PriceDA.Data[2514] := 0.0490536;
   Prof_PriceDA.Data[2515] := 0.0490536;
   Prof_PriceDA.Data[2516] := 0.118098;
   Prof_PriceDA.Data[2517] := 0.118098;
   Prof_PriceDA.Data[2518] := 0.118098;
   Prof_PriceDA.Data[2519] := 0.118098;
   Prof_PriceDA.Data[2520] := 0.1559088;
   Prof_PriceDA.Data[2521] := 0.1559088;
   Prof_PriceDA.Data[2522] := 0.1559088;
   Prof_PriceDA.Data[2523] := 0.1559088;
   Prof_PriceDA.Data[2524] := 0.187002;
   Prof_PriceDA.Data[2525] := 0.187002;
   Prof_PriceDA.Data[2526] := 0.187002;
   Prof_PriceDA.Data[2527] := 0.187002;
   Prof_PriceDA.Data[2528] := 0.1719684;
   Prof_PriceDA.Data[2529] := 0.1719684;
   Prof_PriceDA.Data[2530] := 0.1719684;
   Prof_PriceDA.Data[2531] := 0.1719684;
   Prof_PriceDA.Data[2532] := 0.1409616;
   Prof_PriceDA.Data[2533] := 0.1409616;
   Prof_PriceDA.Data[2534] := 0.1409616;
   Prof_PriceDA.Data[2535] := 0.1409616;
   Prof_PriceDA.Data[2536] := 0.1084428;
   Prof_PriceDA.Data[2537] := 0.1084428;
   Prof_PriceDA.Data[2538] := 0.1084428;
   Prof_PriceDA.Data[2539] := 0.1084428;
   Prof_PriceDA.Data[2540] := 0.1040148;
   Prof_PriceDA.Data[2541] := 0.1040148;
   Prof_PriceDA.Data[2542] := 0.1040148;
   Prof_PriceDA.Data[2543] := 0.1040148;
   Prof_PriceDA.Data[2544] := 0.0946944;
   Prof_PriceDA.Data[2545] := 0.0946944;
   Prof_PriceDA.Data[2546] := 0.0946944;
   Prof_PriceDA.Data[2547] := 0.0946944;
   Prof_PriceDA.Data[2548] := 0.1125792;
   Prof_PriceDA.Data[2549] := 0.1125792;
   Prof_PriceDA.Data[2550] := 0.1125792;
   Prof_PriceDA.Data[2551] := 0.1125792;
   Prof_PriceDA.Data[2552] := 0.1399464;
   Prof_PriceDA.Data[2553] := 0.1399464;
   Prof_PriceDA.Data[2554] := 0.1399464;
   Prof_PriceDA.Data[2555] := 0.1399464;
   Prof_PriceDA.Data[2556] := 0.1582416;
   Prof_PriceDA.Data[2557] := 0.1582416;
   Prof_PriceDA.Data[2558] := 0.1582416;
   Prof_PriceDA.Data[2559] := 0.1582416;
   Prof_PriceDA.Data[2560] := 0.1937628;
   Prof_PriceDA.Data[2561] := 0.1937628;
   Prof_PriceDA.Data[2562] := 0.1937628;
   Prof_PriceDA.Data[2563] := 0.1937628;
   Prof_PriceDA.Data[2564] := 0.1899936;
   Prof_PriceDA.Data[2565] := 0.1899936;
   Prof_PriceDA.Data[2566] := 0.1899936;
   Prof_PriceDA.Data[2567] := 0.1899936;
   Prof_PriceDA.Data[2568] := 0.1928124;
   Prof_PriceDA.Data[2569] := 0.1928124;
   Prof_PriceDA.Data[2570] := 0.1928124;
   Prof_PriceDA.Data[2571] := 0.1928124;
   Prof_PriceDA.Data[2572] := 0.1906308;
   Prof_PriceDA.Data[2573] := 0.1906308;
   Prof_PriceDA.Data[2574] := 0.1906308;
   Prof_PriceDA.Data[2575] := 0.1906308;
   Prof_PriceDA.Data[2576] := 0.170856;
   Prof_PriceDA.Data[2577] := 0.170856;
   Prof_PriceDA.Data[2578] := 0.170856;
   Prof_PriceDA.Data[2579] := 0.170856;
   Prof_PriceDA.Data[2580] := 0.1461024;
   Prof_PriceDA.Data[2581] := 0.1461024;
   Prof_PriceDA.Data[2582] := 0.1461024;
   Prof_PriceDA.Data[2583] := 0.1461024;
   Prof_PriceDA.Data[2584] := 0.130626;
   Prof_PriceDA.Data[2585] := 0.130626;
   Prof_PriceDA.Data[2586] := 0.130626;
   Prof_PriceDA.Data[2587] := 0.130626;
   Prof_PriceDA.Data[2588] := 0.106056;
   Prof_PriceDA.Data[2589] := 0.106056;
   Prof_PriceDA.Data[2590] := 0.106056;
   Prof_PriceDA.Data[2591] := 0.106056;
   Prof_PriceDA.Data[2592] := 0.106758;
   Prof_PriceDA.Data[2593] := 0.106758;
   Prof_PriceDA.Data[2594] := 0.106758;
   Prof_PriceDA.Data[2595] := 0.106758;
   Prof_PriceDA.Data[2596] := 0.0855684;
   Prof_PriceDA.Data[2597] := 0.0855684;
   Prof_PriceDA.Data[2598] := 0.0855684;
   Prof_PriceDA.Data[2599] := 0.0855684;
   Prof_PriceDA.Data[2600] := 0.0941112;
   Prof_PriceDA.Data[2601] := 0.0941112;
   Prof_PriceDA.Data[2602] := 0.0941112;
   Prof_PriceDA.Data[2603] := 0.0941112;
   Prof_PriceDA.Data[2604] := 0.0877068;
   Prof_PriceDA.Data[2605] := 0.0877068;
   Prof_PriceDA.Data[2606] := 0.0877068;
   Prof_PriceDA.Data[2607] := 0.0877068;
   Prof_PriceDA.Data[2608] := 0.0877392;
   Prof_PriceDA.Data[2609] := 0.0877392;
   Prof_PriceDA.Data[2610] := 0.0877392;
   Prof_PriceDA.Data[2611] := 0.0877392;
   Prof_PriceDA.Data[2612] := 0.122688;
   Prof_PriceDA.Data[2613] := 0.122688;
   Prof_PriceDA.Data[2614] := 0.122688;
   Prof_PriceDA.Data[2615] := 0.122688;
   Prof_PriceDA.Data[2616] := 0.1498608;
   Prof_PriceDA.Data[2617] := 0.1498608;
   Prof_PriceDA.Data[2618] := 0.1498608;
   Prof_PriceDA.Data[2619] := 0.1498608;
   Prof_PriceDA.Data[2620] := 0.1502712;
   Prof_PriceDA.Data[2621] := 0.1502712;
   Prof_PriceDA.Data[2622] := 0.1502712;
   Prof_PriceDA.Data[2623] := 0.1502712;
   Prof_PriceDA.Data[2624] := 0.1519992;
   Prof_PriceDA.Data[2625] := 0.1519992;
   Prof_PriceDA.Data[2626] := 0.1519992;
   Prof_PriceDA.Data[2627] := 0.1519992;
   Prof_PriceDA.Data[2628] := 0.1354212;
   Prof_PriceDA.Data[2629] := 0.1354212;
   Prof_PriceDA.Data[2630] := 0.1354212;
   Prof_PriceDA.Data[2631] := 0.1354212;
   Prof_PriceDA.Data[2632] := 0.141318;
   Prof_PriceDA.Data[2633] := 0.141318;
   Prof_PriceDA.Data[2634] := 0.141318;
   Prof_PriceDA.Data[2635] := 0.141318;
   Prof_PriceDA.Data[2636] := 0.1357344;
   Prof_PriceDA.Data[2637] := 0.1357344;
   Prof_PriceDA.Data[2638] := 0.1357344;
   Prof_PriceDA.Data[2639] := 0.1357344;
   Prof_PriceDA.Data[2640] := 0.1322892;
   Prof_PriceDA.Data[2641] := 0.1322892;
   Prof_PriceDA.Data[2642] := 0.1322892;
   Prof_PriceDA.Data[2643] := 0.1322892;
   Prof_PriceDA.Data[2644] := 0.1372788;
   Prof_PriceDA.Data[2645] := 0.1372788;
   Prof_PriceDA.Data[2646] := 0.1372788;
   Prof_PriceDA.Data[2647] := 0.1372788;
   Prof_PriceDA.Data[2648] := 0.1420632;
   Prof_PriceDA.Data[2649] := 0.1420632;
   Prof_PriceDA.Data[2650] := 0.1420632;
   Prof_PriceDA.Data[2651] := 0.1420632;
   Prof_PriceDA.Data[2652] := 0.135162;
   Prof_PriceDA.Data[2653] := 0.135162;
   Prof_PriceDA.Data[2654] := 0.135162;
   Prof_PriceDA.Data[2655] := 0.135162;
   Prof_PriceDA.Data[2656] := 0.1540296;
   Prof_PriceDA.Data[2657] := 0.1540296;
   Prof_PriceDA.Data[2658] := 0.1540296;
   Prof_PriceDA.Data[2659] := 0.1540296;
   Prof_PriceDA.Data[2660] := 0.1559304;
   Prof_PriceDA.Data[2661] := 0.1559304;
   Prof_PriceDA.Data[2662] := 0.1559304;
   Prof_PriceDA.Data[2663] := 0.1559304;
   Prof_PriceDA.Data[2664] := 0.1593864;
   Prof_PriceDA.Data[2665] := 0.1593864;
   Prof_PriceDA.Data[2666] := 0.1593864;
   Prof_PriceDA.Data[2667] := 0.1593864;
   Prof_PriceDA.Data[2668] := 0.1502928;
   Prof_PriceDA.Data[2669] := 0.1502928;
   Prof_PriceDA.Data[2670] := 0.1502928;
   Prof_PriceDA.Data[2671] := 0.1502928;
   Prof_PriceDA.Data[2672] := 0.1499256;
   Prof_PriceDA.Data[2673] := 0.1499256;
   Prof_PriceDA.Data[2674] := 0.1499256;
   Prof_PriceDA.Data[2675] := 0.1499256;
   Prof_PriceDA.Data[2676] := 0.1251612;
   Prof_PriceDA.Data[2677] := 0.1251612;
   Prof_PriceDA.Data[2678] := 0.1251612;
   Prof_PriceDA.Data[2679] := 0.1251612;
   Prof_PriceDA.Data[2680] := 0.1250208;
   Prof_PriceDA.Data[2681] := 0.1250208;
   Prof_PriceDA.Data[2682] := 0.1250208;
   Prof_PriceDA.Data[2683] := 0.1250208;
   Prof_PriceDA.Data[2684] := 0.1051704;
   Prof_PriceDA.Data[2685] := 0.1051704;
   Prof_PriceDA.Data[2686] := 0.1051704;
   Prof_PriceDA.Data[2687] := 0.1051704;
   Prof_PriceDA.Data[2688] := 0.105462;
   Prof_PriceDA.Data[2689] := 0.105462;
   Prof_PriceDA.Data[2690] := 0.105462;
   Prof_PriceDA.Data[2691] := 0.105462;
   Prof_PriceDA.Data[2692] := 0.097362;
   Prof_PriceDA.Data[2693] := 0.097362;
   Prof_PriceDA.Data[2694] := 0.097362;
   Prof_PriceDA.Data[2695] := 0.097362;
   Prof_PriceDA.Data[2696] := 0.0910332;
   Prof_PriceDA.Data[2697] := 0.0910332;
   Prof_PriceDA.Data[2698] := 0.0910332;
   Prof_PriceDA.Data[2699] := 0.0910332;
   Prof_PriceDA.Data[2700] := 0.0914328;
   Prof_PriceDA.Data[2701] := 0.0914328;
   Prof_PriceDA.Data[2702] := 0.0914328;
   Prof_PriceDA.Data[2703] := 0.0914328;
   Prof_PriceDA.Data[2704] := 0.0972;
   Prof_PriceDA.Data[2705] := 0.0972;
   Prof_PriceDA.Data[2706] := 0.0972;
   Prof_PriceDA.Data[2707] := 0.0972;
   Prof_PriceDA.Data[2708] := 0.1214676;
   Prof_PriceDA.Data[2709] := 0.1214676;
   Prof_PriceDA.Data[2710] := 0.1214676;
   Prof_PriceDA.Data[2711] := 0.1214676;
   Prof_PriceDA.Data[2712] := 0.154656;
   Prof_PriceDA.Data[2713] := 0.154656;
   Prof_PriceDA.Data[2714] := 0.154656;
   Prof_PriceDA.Data[2715] := 0.154656;
   Prof_PriceDA.Data[2716] := 0.1773468;
   Prof_PriceDA.Data[2717] := 0.1773468;
   Prof_PriceDA.Data[2718] := 0.1773468;
   Prof_PriceDA.Data[2719] := 0.1773468;
   Prof_PriceDA.Data[2720] := 0.1579068;
   Prof_PriceDA.Data[2721] := 0.1579068;
   Prof_PriceDA.Data[2722] := 0.1579068;
   Prof_PriceDA.Data[2723] := 0.1579068;
   Prof_PriceDA.Data[2724] := 0.1480896;
   Prof_PriceDA.Data[2725] := 0.1480896;
   Prof_PriceDA.Data[2726] := 0.1480896;
   Prof_PriceDA.Data[2727] := 0.1480896;
   Prof_PriceDA.Data[2728] := 0.1204308;
   Prof_PriceDA.Data[2729] := 0.1204308;
   Prof_PriceDA.Data[2730] := 0.1204308;
   Prof_PriceDA.Data[2731] := 0.1204308;
   Prof_PriceDA.Data[2732] := 0.1014444;
   Prof_PriceDA.Data[2733] := 0.1014444;
   Prof_PriceDA.Data[2734] := 0.1014444;
   Prof_PriceDA.Data[2735] := 0.1014444;
   Prof_PriceDA.Data[2736] := 0.093204;
   Prof_PriceDA.Data[2737] := 0.093204;
   Prof_PriceDA.Data[2738] := 0.093204;
   Prof_PriceDA.Data[2739] := 0.093204;
   Prof_PriceDA.Data[2740] := 0.0935496;
   Prof_PriceDA.Data[2741] := 0.0935496;
   Prof_PriceDA.Data[2742] := 0.0935496;
   Prof_PriceDA.Data[2743] := 0.0935496;
   Prof_PriceDA.Data[2744] := 0.1055484;
   Prof_PriceDA.Data[2745] := 0.1055484;
   Prof_PriceDA.Data[2746] := 0.1055484;
   Prof_PriceDA.Data[2747] := 0.1055484;
   Prof_PriceDA.Data[2748] := 0.1400328;
   Prof_PriceDA.Data[2749] := 0.1400328;
   Prof_PriceDA.Data[2750] := 0.1400328;
   Prof_PriceDA.Data[2751] := 0.1400328;
   Prof_PriceDA.Data[2752] := 0.1792692;
   Prof_PriceDA.Data[2753] := 0.1792692;
   Prof_PriceDA.Data[2754] := 0.1792692;
   Prof_PriceDA.Data[2755] := 0.1792692;
   Prof_PriceDA.Data[2756] := 0.1827792;
   Prof_PriceDA.Data[2757] := 0.1827792;
   Prof_PriceDA.Data[2758] := 0.1827792;
   Prof_PriceDA.Data[2759] := 0.1827792;
   Prof_PriceDA.Data[2760] := 0.1721088;
   Prof_PriceDA.Data[2761] := 0.1721088;
   Prof_PriceDA.Data[2762] := 0.1721088;
   Prof_PriceDA.Data[2763] := 0.1721088;
   Prof_PriceDA.Data[2764] := 0.173502;
   Prof_PriceDA.Data[2765] := 0.173502;
   Prof_PriceDA.Data[2766] := 0.173502;
   Prof_PriceDA.Data[2767] := 0.173502;
   Prof_PriceDA.Data[2768] := 0.1609524;
   Prof_PriceDA.Data[2769] := 0.1609524;
   Prof_PriceDA.Data[2770] := 0.1609524;
   Prof_PriceDA.Data[2771] := 0.1609524;
   Prof_PriceDA.Data[2772] := 0.1491912;
   Prof_PriceDA.Data[2773] := 0.1491912;
   Prof_PriceDA.Data[2774] := 0.1491912;
   Prof_PriceDA.Data[2775] := 0.1491912;
   Prof_PriceDA.Data[2776] := 0.1330236;
   Prof_PriceDA.Data[2777] := 0.1330236;
   Prof_PriceDA.Data[2778] := 0.1330236;
   Prof_PriceDA.Data[2779] := 0.1330236;
   Prof_PriceDA.Data[2780] := 0.1119204;
   Prof_PriceDA.Data[2781] := 0.1119204;
   Prof_PriceDA.Data[2782] := 0.1119204;
   Prof_PriceDA.Data[2783] := 0.1119204;
   Prof_PriceDA.Data[2784] := 0.110268;
   Prof_PriceDA.Data[2785] := 0.110268;
   Prof_PriceDA.Data[2786] := 0.110268;
   Prof_PriceDA.Data[2787] := 0.110268;
   Prof_PriceDA.Data[2788] := 0.1095228;
   Prof_PriceDA.Data[2789] := 0.1095228;
   Prof_PriceDA.Data[2790] := 0.1095228;
   Prof_PriceDA.Data[2791] := 0.1095228;
   Prof_PriceDA.Data[2792] := 0.1069524;
   Prof_PriceDA.Data[2793] := 0.1069524;
   Prof_PriceDA.Data[2794] := 0.1069524;
   Prof_PriceDA.Data[2795] := 0.1069524;
   Prof_PriceDA.Data[2796] := 0.1100844;
   Prof_PriceDA.Data[2797] := 0.1100844;
   Prof_PriceDA.Data[2798] := 0.1100844;
   Prof_PriceDA.Data[2799] := 0.1100844;
   Prof_PriceDA.Data[2800] := 0.1098036;
   Prof_PriceDA.Data[2801] := 0.1098036;
   Prof_PriceDA.Data[2802] := 0.1098036;
   Prof_PriceDA.Data[2803] := 0.1098036;
   Prof_PriceDA.Data[2804] := 0.1232496;
   Prof_PriceDA.Data[2805] := 0.1232496;
   Prof_PriceDA.Data[2806] := 0.1232496;
   Prof_PriceDA.Data[2807] := 0.1232496;
   Prof_PriceDA.Data[2808] := 0.1569348;
   Prof_PriceDA.Data[2809] := 0.1569348;
   Prof_PriceDA.Data[2810] := 0.1569348;
   Prof_PriceDA.Data[2811] := 0.1569348;
   Prof_PriceDA.Data[2812] := 0.1669788;
   Prof_PriceDA.Data[2813] := 0.1669788;
   Prof_PriceDA.Data[2814] := 0.1669788;
   Prof_PriceDA.Data[2815] := 0.1669788;
   Prof_PriceDA.Data[2816] := 0.173124;
   Prof_PriceDA.Data[2817] := 0.173124;
   Prof_PriceDA.Data[2818] := 0.173124;
   Prof_PriceDA.Data[2819] := 0.173124;
   Prof_PriceDA.Data[2820] := 0.1639764;
   Prof_PriceDA.Data[2821] := 0.1639764;
   Prof_PriceDA.Data[2822] := 0.1639764;
   Prof_PriceDA.Data[2823] := 0.1639764;
   Prof_PriceDA.Data[2824] := 0.1429704;
   Prof_PriceDA.Data[2825] := 0.1429704;
   Prof_PriceDA.Data[2826] := 0.1429704;
   Prof_PriceDA.Data[2827] := 0.1429704;
   Prof_PriceDA.Data[2828] := 0.13311;
   Prof_PriceDA.Data[2829] := 0.13311;
   Prof_PriceDA.Data[2830] := 0.13311;
   Prof_PriceDA.Data[2831] := 0.13311;
   Prof_PriceDA.Data[2832] := 0.1219428;
   Prof_PriceDA.Data[2833] := 0.1219428;
   Prof_PriceDA.Data[2834] := 0.1219428;
   Prof_PriceDA.Data[2835] := 0.1219428;
   Prof_PriceDA.Data[2836] := 0.122364;
   Prof_PriceDA.Data[2837] := 0.122364;
   Prof_PriceDA.Data[2838] := 0.122364;
   Prof_PriceDA.Data[2839] := 0.122364;
   Prof_PriceDA.Data[2840] := 0.1403892;
   Prof_PriceDA.Data[2841] := 0.1403892;
   Prof_PriceDA.Data[2842] := 0.1403892;
   Prof_PriceDA.Data[2843] := 0.1403892;
   Prof_PriceDA.Data[2844] := 0.1655748;
   Prof_PriceDA.Data[2845] := 0.1655748;
   Prof_PriceDA.Data[2846] := 0.1655748;
   Prof_PriceDA.Data[2847] := 0.1655748;
   Prof_PriceDA.Data[2848] := 0.1736748;
   Prof_PriceDA.Data[2849] := 0.1736748;
   Prof_PriceDA.Data[2850] := 0.1736748;
   Prof_PriceDA.Data[2851] := 0.1736748;
   Prof_PriceDA.Data[2852] := 0.1896696;
   Prof_PriceDA.Data[2853] := 0.1896696;
   Prof_PriceDA.Data[2854] := 0.1896696;
   Prof_PriceDA.Data[2855] := 0.1896696;
   Prof_PriceDA.Data[2856] := 0.1858032;
   Prof_PriceDA.Data[2857] := 0.1858032;
   Prof_PriceDA.Data[2858] := 0.1858032;
   Prof_PriceDA.Data[2859] := 0.1858032;
   Prof_PriceDA.Data[2860] := 0.1741824;
   Prof_PriceDA.Data[2861] := 0.1741824;
   Prof_PriceDA.Data[2862] := 0.1741824;
   Prof_PriceDA.Data[2863] := 0.1741824;
   Prof_PriceDA.Data[2864] := 0.1635228;
   Prof_PriceDA.Data[2865] := 0.1635228;
   Prof_PriceDA.Data[2866] := 0.1635228;
   Prof_PriceDA.Data[2867] := 0.1635228;
   Prof_PriceDA.Data[2868] := 0.145908;
   Prof_PriceDA.Data[2869] := 0.145908;
   Prof_PriceDA.Data[2870] := 0.145908;
   Prof_PriceDA.Data[2871] := 0.145908;
   Prof_PriceDA.Data[2872] := 0.1370952;
   Prof_PriceDA.Data[2873] := 0.1370952;
   Prof_PriceDA.Data[2874] := 0.1370952;
   Prof_PriceDA.Data[2875] := 0.1370952;
   Prof_PriceDA.Data[2876] := 0.129816;
   Prof_PriceDA.Data[2877] := 0.129816;
   Prof_PriceDA.Data[2878] := 0.129816;
   Prof_PriceDA.Data[2879] := 0.129816;
   Prof_PriceDA.Data[2880] := 0.1296;
   Prof_PriceDA.Data[2881] := 0.1296;
   Prof_PriceDA.Data[2882] := 0.1296;
   Prof_PriceDA.Data[2883] := 0.1296;
   Prof_PriceDA.Data[2884] := 0.1269;
   Prof_PriceDA.Data[2885] := 0.1269;
   Prof_PriceDA.Data[2886] := 0.1269;
   Prof_PriceDA.Data[2887] := 0.1269;
   Prof_PriceDA.Data[2888] := 0.1232064;
   Prof_PriceDA.Data[2889] := 0.1232064;
   Prof_PriceDA.Data[2890] := 0.1232064;
   Prof_PriceDA.Data[2891] := 0.1232064;
   Prof_PriceDA.Data[2892] := 0.1236384;
   Prof_PriceDA.Data[2893] := 0.1236384;
   Prof_PriceDA.Data[2894] := 0.1236384;
   Prof_PriceDA.Data[2895] := 0.1236384;
   Prof_PriceDA.Data[2896] := 0.1267164;
   Prof_PriceDA.Data[2897] := 0.1267164;
   Prof_PriceDA.Data[2898] := 0.1267164;
   Prof_PriceDA.Data[2899] := 0.1267164;
   Prof_PriceDA.Data[2900] := 0.1316088;
   Prof_PriceDA.Data[2901] := 0.1316088;
   Prof_PriceDA.Data[2902] := 0.1316088;
   Prof_PriceDA.Data[2903] := 0.1316088;
   Prof_PriceDA.Data[2904] := 0.1604556;
   Prof_PriceDA.Data[2905] := 0.1604556;
   Prof_PriceDA.Data[2906] := 0.1604556;
   Prof_PriceDA.Data[2907] := 0.1604556;
   Prof_PriceDA.Data[2908] := 0.1728;
   Prof_PriceDA.Data[2909] := 0.1728;
   Prof_PriceDA.Data[2910] := 0.1728;
   Prof_PriceDA.Data[2911] := 0.1728;
   Prof_PriceDA.Data[2912] := 0.176796;
   Prof_PriceDA.Data[2913] := 0.176796;
   Prof_PriceDA.Data[2914] := 0.176796;
   Prof_PriceDA.Data[2915] := 0.176796;
   Prof_PriceDA.Data[2916] := 0.1672056;
   Prof_PriceDA.Data[2917] := 0.1672056;
   Prof_PriceDA.Data[2918] := 0.1672056;
   Prof_PriceDA.Data[2919] := 0.1672056;
   Prof_PriceDA.Data[2920] := 0.140508;
   Prof_PriceDA.Data[2921] := 0.140508;
   Prof_PriceDA.Data[2922] := 0.140508;
   Prof_PriceDA.Data[2923] := 0.140508;
   Prof_PriceDA.Data[2924] := 0.136296;
   Prof_PriceDA.Data[2925] := 0.136296;
   Prof_PriceDA.Data[2926] := 0.136296;
   Prof_PriceDA.Data[2927] := 0.136296;
   Prof_PriceDA.Data[2928] := 0.1296648;
   Prof_PriceDA.Data[2929] := 0.1296648;
   Prof_PriceDA.Data[2930] := 0.1296648;
   Prof_PriceDA.Data[2931] := 0.1296648;
   Prof_PriceDA.Data[2932] := 0.1308852;
   Prof_PriceDA.Data[2933] := 0.1308852;
   Prof_PriceDA.Data[2934] := 0.1308852;
   Prof_PriceDA.Data[2935] := 0.1308852;
   Prof_PriceDA.Data[2936] := 0.1296432;
   Prof_PriceDA.Data[2937] := 0.1296432;
   Prof_PriceDA.Data[2938] := 0.1296432;
   Prof_PriceDA.Data[2939] := 0.1296432;
   Prof_PriceDA.Data[2940] := 0.1655964;
   Prof_PriceDA.Data[2941] := 0.1655964;
   Prof_PriceDA.Data[2942] := 0.1655964;
   Prof_PriceDA.Data[2943] := 0.1655964;
   Prof_PriceDA.Data[2944] := 0.1810512;
   Prof_PriceDA.Data[2945] := 0.1810512;
   Prof_PriceDA.Data[2946] := 0.1810512;
   Prof_PriceDA.Data[2947] := 0.1810512;
   Prof_PriceDA.Data[2948] := 0.1930716;
   Prof_PriceDA.Data[2949] := 0.1930716;
   Prof_PriceDA.Data[2950] := 0.1930716;
   Prof_PriceDA.Data[2951] := 0.1930716;
   Prof_PriceDA.Data[2952] := 0.1992384;
   Prof_PriceDA.Data[2953] := 0.1992384;
   Prof_PriceDA.Data[2954] := 0.1992384;
   Prof_PriceDA.Data[2955] := 0.1992384;
   Prof_PriceDA.Data[2956] := 0.1933092;
   Prof_PriceDA.Data[2957] := 0.1933092;
   Prof_PriceDA.Data[2958] := 0.1933092;
   Prof_PriceDA.Data[2959] := 0.1933092;
   Prof_PriceDA.Data[2960] := 0.1756728;
   Prof_PriceDA.Data[2961] := 0.1756728;
   Prof_PriceDA.Data[2962] := 0.1756728;
   Prof_PriceDA.Data[2963] := 0.1756728;
   Prof_PriceDA.Data[2964] := 0.164916;
   Prof_PriceDA.Data[2965] := 0.164916;
   Prof_PriceDA.Data[2966] := 0.164916;
   Prof_PriceDA.Data[2967] := 0.164916;
   Prof_PriceDA.Data[2968] := 0.1607472;
   Prof_PriceDA.Data[2969] := 0.1607472;
   Prof_PriceDA.Data[2970] := 0.1607472;
   Prof_PriceDA.Data[2971] := 0.1607472;
   Prof_PriceDA.Data[2972] := 0.144126;
   Prof_PriceDA.Data[2973] := 0.144126;
   Prof_PriceDA.Data[2974] := 0.144126;
   Prof_PriceDA.Data[2975] := 0.144126;
   Prof_PriceDA.Data[2976] := 0.1494828;
   Prof_PriceDA.Data[2977] := 0.1494828;
   Prof_PriceDA.Data[2978] := 0.1494828;
   Prof_PriceDA.Data[2979] := 0.1494828;
   Prof_PriceDA.Data[2980] := 0.1409724;
   Prof_PriceDA.Data[2981] := 0.1409724;
   Prof_PriceDA.Data[2982] := 0.1409724;
   Prof_PriceDA.Data[2983] := 0.1409724;
   Prof_PriceDA.Data[2984] := 0.135108;
   Prof_PriceDA.Data[2985] := 0.135108;
   Prof_PriceDA.Data[2986] := 0.135108;
   Prof_PriceDA.Data[2987] := 0.135108;
   Prof_PriceDA.Data[2988] := 0.1288332;
   Prof_PriceDA.Data[2989] := 0.1288332;
   Prof_PriceDA.Data[2990] := 0.1288332;
   Prof_PriceDA.Data[2991] := 0.1288332;
   Prof_PriceDA.Data[2992] := 0.1295568;
   Prof_PriceDA.Data[2993] := 0.1295568;
   Prof_PriceDA.Data[2994] := 0.1295568;
   Prof_PriceDA.Data[2995] := 0.1295568;
   Prof_PriceDA.Data[2996] := 0.1312308;
   Prof_PriceDA.Data[2997] := 0.1312308;
   Prof_PriceDA.Data[2998] := 0.1312308;
   Prof_PriceDA.Data[2999] := 0.1312308;
   Prof_PriceDA.Data[3000] := 0.1374948;
   Prof_PriceDA.Data[3001] := 0.1374948;
   Prof_PriceDA.Data[3002] := 0.1374948;
   Prof_PriceDA.Data[3003] := 0.1374948;
   Prof_PriceDA.Data[3004] := 0.1563192;
   Prof_PriceDA.Data[3005] := 0.1563192;
   Prof_PriceDA.Data[3006] := 0.1563192;
   Prof_PriceDA.Data[3007] := 0.1563192;
   Prof_PriceDA.Data[3008] := 0.1657368;
   Prof_PriceDA.Data[3009] := 0.1657368;
   Prof_PriceDA.Data[3010] := 0.1657368;
   Prof_PriceDA.Data[3011] := 0.1657368;
   Prof_PriceDA.Data[3012] := 0.1538352;
   Prof_PriceDA.Data[3013] := 0.1538352;
   Prof_PriceDA.Data[3014] := 0.1538352;
   Prof_PriceDA.Data[3015] := 0.1538352;
   Prof_PriceDA.Data[3016] := 0.138672;
   Prof_PriceDA.Data[3017] := 0.138672;
   Prof_PriceDA.Data[3018] := 0.138672;
   Prof_PriceDA.Data[3019] := 0.138672;
   Prof_PriceDA.Data[3020] := 0.1296864;
   Prof_PriceDA.Data[3021] := 0.1296864;
   Prof_PriceDA.Data[3022] := 0.1296864;
   Prof_PriceDA.Data[3023] := 0.1296864;
   Prof_PriceDA.Data[3024] := 0.1191132;
   Prof_PriceDA.Data[3025] := 0.1191132;
   Prof_PriceDA.Data[3026] := 0.1191132;
   Prof_PriceDA.Data[3027] := 0.1191132;
   Prof_PriceDA.Data[3028] := 0.111672;
   Prof_PriceDA.Data[3029] := 0.111672;
   Prof_PriceDA.Data[3030] := 0.111672;
   Prof_PriceDA.Data[3031] := 0.111672;
   Prof_PriceDA.Data[3032] := 0.122796;
   Prof_PriceDA.Data[3033] := 0.122796;
   Prof_PriceDA.Data[3034] := 0.122796;
   Prof_PriceDA.Data[3035] := 0.122796;
   Prof_PriceDA.Data[3036] := 0.1411344;
   Prof_PriceDA.Data[3037] := 0.1411344;
   Prof_PriceDA.Data[3038] := 0.1411344;
   Prof_PriceDA.Data[3039] := 0.1411344;
   Prof_PriceDA.Data[3040] := 0.1683072;
   Prof_PriceDA.Data[3041] := 0.1683072;
   Prof_PriceDA.Data[3042] := 0.1683072;
   Prof_PriceDA.Data[3043] := 0.1683072;
   Prof_PriceDA.Data[3044] := 0.1792368;
   Prof_PriceDA.Data[3045] := 0.1792368;
   Prof_PriceDA.Data[3046] := 0.1792368;
   Prof_PriceDA.Data[3047] := 0.1792368;
   Prof_PriceDA.Data[3048] := 0.180036;
   Prof_PriceDA.Data[3049] := 0.180036;
   Prof_PriceDA.Data[3050] := 0.180036;
   Prof_PriceDA.Data[3051] := 0.180036;
   Prof_PriceDA.Data[3052] := 0.1760184;
   Prof_PriceDA.Data[3053] := 0.1760184;
   Prof_PriceDA.Data[3054] := 0.1760184;
   Prof_PriceDA.Data[3055] := 0.1760184;
   Prof_PriceDA.Data[3056] := 0.169128;
   Prof_PriceDA.Data[3057] := 0.169128;
   Prof_PriceDA.Data[3058] := 0.169128;
   Prof_PriceDA.Data[3059] := 0.169128;
   Prof_PriceDA.Data[3060] := 0.1568592;
   Prof_PriceDA.Data[3061] := 0.1568592;
   Prof_PriceDA.Data[3062] := 0.1568592;
   Prof_PriceDA.Data[3063] := 0.1568592;
   Prof_PriceDA.Data[3064] := 0.1530684;
   Prof_PriceDA.Data[3065] := 0.1530684;
   Prof_PriceDA.Data[3066] := 0.1530684;
   Prof_PriceDA.Data[3067] := 0.1530684;
   Prof_PriceDA.Data[3068] := 0.1422792;
   Prof_PriceDA.Data[3069] := 0.1422792;
   Prof_PriceDA.Data[3070] := 0.1422792;
   Prof_PriceDA.Data[3071] := 0.1422792;
   Prof_PriceDA.Data[3072] := 0.1439208;
   Prof_PriceDA.Data[3073] := 0.1439208;
   Prof_PriceDA.Data[3074] := 0.1439208;
   Prof_PriceDA.Data[3075] := 0.1439208;
   Prof_PriceDA.Data[3076] := 0.1370628;
   Prof_PriceDA.Data[3077] := 0.1370628;
   Prof_PriceDA.Data[3078] := 0.1370628;
   Prof_PriceDA.Data[3079] := 0.1370628;
   Prof_PriceDA.Data[3080] := 0.1328292;
   Prof_PriceDA.Data[3081] := 0.1328292;
   Prof_PriceDA.Data[3082] := 0.1328292;
   Prof_PriceDA.Data[3083] := 0.1328292;
   Prof_PriceDA.Data[3084] := 0.1303128;
   Prof_PriceDA.Data[3085] := 0.1303128;
   Prof_PriceDA.Data[3086] := 0.1303128;
   Prof_PriceDA.Data[3087] := 0.1303128;
   Prof_PriceDA.Data[3088] := 0.1321272;
   Prof_PriceDA.Data[3089] := 0.1321272;
   Prof_PriceDA.Data[3090] := 0.1321272;
   Prof_PriceDA.Data[3091] := 0.1321272;
   Prof_PriceDA.Data[3092] := 0.1332828;
   Prof_PriceDA.Data[3093] := 0.1332828;
   Prof_PriceDA.Data[3094] := 0.1332828;
   Prof_PriceDA.Data[3095] := 0.1332828;
   Prof_PriceDA.Data[3096] := 0.1383372;
   Prof_PriceDA.Data[3097] := 0.1383372;
   Prof_PriceDA.Data[3098] := 0.1383372;
   Prof_PriceDA.Data[3099] := 0.1383372;
   Prof_PriceDA.Data[3100] := 0.146772;
   Prof_PriceDA.Data[3101] := 0.146772;
   Prof_PriceDA.Data[3102] := 0.146772;
   Prof_PriceDA.Data[3103] := 0.146772;
   Prof_PriceDA.Data[3104] := 0.148284;
   Prof_PriceDA.Data[3105] := 0.148284;
   Prof_PriceDA.Data[3106] := 0.148284;
   Prof_PriceDA.Data[3107] := 0.148284;
   Prof_PriceDA.Data[3108] := 0.148716;
   Prof_PriceDA.Data[3109] := 0.148716;
   Prof_PriceDA.Data[3110] := 0.148716;
   Prof_PriceDA.Data[3111] := 0.148716;
   Prof_PriceDA.Data[3112] := 0.1404432;
   Prof_PriceDA.Data[3113] := 0.1404432;
   Prof_PriceDA.Data[3114] := 0.1404432;
   Prof_PriceDA.Data[3115] := 0.1404432;
   Prof_PriceDA.Data[3116] := 0.1396764;
   Prof_PriceDA.Data[3117] := 0.1396764;
   Prof_PriceDA.Data[3118] := 0.1396764;
   Prof_PriceDA.Data[3119] := 0.1396764;
   Prof_PriceDA.Data[3120] := 0.1320192;
   Prof_PriceDA.Data[3121] := 0.1320192;
   Prof_PriceDA.Data[3122] := 0.1320192;
   Prof_PriceDA.Data[3123] := 0.1320192;
   Prof_PriceDA.Data[3124] := 0.1208304;
   Prof_PriceDA.Data[3125] := 0.1208304;
   Prof_PriceDA.Data[3126] := 0.1208304;
   Prof_PriceDA.Data[3127] := 0.1208304;
   Prof_PriceDA.Data[3128] := 0.1263168;
   Prof_PriceDA.Data[3129] := 0.1263168;
   Prof_PriceDA.Data[3130] := 0.1263168;
   Prof_PriceDA.Data[3131] := 0.1263168;
   Prof_PriceDA.Data[3132] := 0.140562;
   Prof_PriceDA.Data[3133] := 0.140562;
   Prof_PriceDA.Data[3134] := 0.140562;
   Prof_PriceDA.Data[3135] := 0.140562;
   Prof_PriceDA.Data[3136] := 0.168156;
   Prof_PriceDA.Data[3137] := 0.168156;
   Prof_PriceDA.Data[3138] := 0.168156;
   Prof_PriceDA.Data[3139] := 0.168156;
   Prof_PriceDA.Data[3140] := 0.1802088;
   Prof_PriceDA.Data[3141] := 0.1802088;
   Prof_PriceDA.Data[3142] := 0.1802088;
   Prof_PriceDA.Data[3143] := 0.1802088;
   Prof_PriceDA.Data[3144] := 0.185544;
   Prof_PriceDA.Data[3145] := 0.185544;
   Prof_PriceDA.Data[3146] := 0.185544;
   Prof_PriceDA.Data[3147] := 0.185544;
   Prof_PriceDA.Data[3148] := 0.187866;
   Prof_PriceDA.Data[3149] := 0.187866;
   Prof_PriceDA.Data[3150] := 0.187866;
   Prof_PriceDA.Data[3151] := 0.187866;
   Prof_PriceDA.Data[3152] := 0.17874;
   Prof_PriceDA.Data[3153] := 0.17874;
   Prof_PriceDA.Data[3154] := 0.17874;
   Prof_PriceDA.Data[3155] := 0.17874;
   Prof_PriceDA.Data[3156] := 0.1682316;
   Prof_PriceDA.Data[3157] := 0.1682316;
   Prof_PriceDA.Data[3158] := 0.1682316;
   Prof_PriceDA.Data[3159] := 0.1682316;
   Prof_PriceDA.Data[3160] := 0.1603152;
   Prof_PriceDA.Data[3161] := 0.1603152;
   Prof_PriceDA.Data[3162] := 0.1603152;
   Prof_PriceDA.Data[3163] := 0.1603152;
   Prof_PriceDA.Data[3164] := 0.1438992;
   Prof_PriceDA.Data[3165] := 0.1438992;
   Prof_PriceDA.Data[3166] := 0.1438992;
   Prof_PriceDA.Data[3167] := 0.1438992;
   Prof_PriceDA.Data[3168] := 0.1399032;
   Prof_PriceDA.Data[3169] := 0.1399032;
   Prof_PriceDA.Data[3170] := 0.1399032;
   Prof_PriceDA.Data[3171] := 0.1399032;
   Prof_PriceDA.Data[3172] := 0.1367604;
   Prof_PriceDA.Data[3173] := 0.1367604;
   Prof_PriceDA.Data[3174] := 0.1367604;
   Prof_PriceDA.Data[3175] := 0.1367604;
   Prof_PriceDA.Data[3176] := 0.1346976;
   Prof_PriceDA.Data[3177] := 0.1346976;
   Prof_PriceDA.Data[3178] := 0.1346976;
   Prof_PriceDA.Data[3179] := 0.1346976;
   Prof_PriceDA.Data[3180] := 0.1296432;
   Prof_PriceDA.Data[3181] := 0.1296432;
   Prof_PriceDA.Data[3182] := 0.1296432;
   Prof_PriceDA.Data[3183] := 0.1296432;
   Prof_PriceDA.Data[3184] := 0.1330992;
   Prof_PriceDA.Data[3185] := 0.1330992;
   Prof_PriceDA.Data[3186] := 0.1330992;
   Prof_PriceDA.Data[3187] := 0.1330992;
   Prof_PriceDA.Data[3188] := 0.1379916;
   Prof_PriceDA.Data[3189] := 0.1379916;
   Prof_PriceDA.Data[3190] := 0.1379916;
   Prof_PriceDA.Data[3191] := 0.1379916;
   Prof_PriceDA.Data[3192] := 0.1719144;
   Prof_PriceDA.Data[3193] := 0.1719144;
   Prof_PriceDA.Data[3194] := 0.1719144;
   Prof_PriceDA.Data[3195] := 0.1719144;
   Prof_PriceDA.Data[3196] := 0.2245104;
   Prof_PriceDA.Data[3197] := 0.2245104;
   Prof_PriceDA.Data[3198] := 0.2245104;
   Prof_PriceDA.Data[3199] := 0.2245104;
   Prof_PriceDA.Data[3200] := 0.2626884;
   Prof_PriceDA.Data[3201] := 0.2626884;
   Prof_PriceDA.Data[3202] := 0.2626884;
   Prof_PriceDA.Data[3203] := 0.2626884;
   Prof_PriceDA.Data[3204] := 0.1922832;
   Prof_PriceDA.Data[3205] := 0.1922832;
   Prof_PriceDA.Data[3206] := 0.1922832;
   Prof_PriceDA.Data[3207] := 0.1922832;
   Prof_PriceDA.Data[3208] := 0.161946;
   Prof_PriceDA.Data[3209] := 0.161946;
   Prof_PriceDA.Data[3210] := 0.161946;
   Prof_PriceDA.Data[3211] := 0.161946;
   Prof_PriceDA.Data[3212] := 0.1363176;
   Prof_PriceDA.Data[3213] := 0.1363176;
   Prof_PriceDA.Data[3214] := 0.1363176;
   Prof_PriceDA.Data[3215] := 0.1363176;
   Prof_PriceDA.Data[3216] := 0.1266516;
   Prof_PriceDA.Data[3217] := 0.1266516;
   Prof_PriceDA.Data[3218] := 0.1266516;
   Prof_PriceDA.Data[3219] := 0.1266516;
   Prof_PriceDA.Data[3220] := 0.1249776;
   Prof_PriceDA.Data[3221] := 0.1249776;
   Prof_PriceDA.Data[3222] := 0.1249776;
   Prof_PriceDA.Data[3223] := 0.1249776;
   Prof_PriceDA.Data[3224] := 0.1344276;
   Prof_PriceDA.Data[3225] := 0.1344276;
   Prof_PriceDA.Data[3226] := 0.1344276;
   Prof_PriceDA.Data[3227] := 0.1344276;
   Prof_PriceDA.Data[3228] := 0.1597968;
   Prof_PriceDA.Data[3229] := 0.1597968;
   Prof_PriceDA.Data[3230] := 0.1597968;
   Prof_PriceDA.Data[3231] := 0.1597968;
   Prof_PriceDA.Data[3232] := 0.1793664;
   Prof_PriceDA.Data[3233] := 0.1793664;
   Prof_PriceDA.Data[3234] := 0.1793664;
   Prof_PriceDA.Data[3235] := 0.1793664;
   Prof_PriceDA.Data[3236] := 0.226962;
   Prof_PriceDA.Data[3237] := 0.226962;
   Prof_PriceDA.Data[3238] := 0.226962;
   Prof_PriceDA.Data[3239] := 0.226962;
   Prof_PriceDA.Data[3240] := 0.2167884;
   Prof_PriceDA.Data[3241] := 0.2167884;
   Prof_PriceDA.Data[3242] := 0.2167884;
   Prof_PriceDA.Data[3243] := 0.2167884;
   Prof_PriceDA.Data[3244] := 0.217188;
   Prof_PriceDA.Data[3245] := 0.217188;
   Prof_PriceDA.Data[3246] := 0.217188;
   Prof_PriceDA.Data[3247] := 0.217188;
   Prof_PriceDA.Data[3248] := 0.1811592;
   Prof_PriceDA.Data[3249] := 0.1811592;
   Prof_PriceDA.Data[3250] := 0.1811592;
   Prof_PriceDA.Data[3251] := 0.1811592;
   Prof_PriceDA.Data[3252] := 0.16524;
   Prof_PriceDA.Data[3253] := 0.16524;
   Prof_PriceDA.Data[3254] := 0.16524;
   Prof_PriceDA.Data[3255] := 0.16524;
   Prof_PriceDA.Data[3256] := 0.1557252;
   Prof_PriceDA.Data[3257] := 0.1557252;
   Prof_PriceDA.Data[3258] := 0.1557252;
   Prof_PriceDA.Data[3259] := 0.1557252;
   Prof_PriceDA.Data[3260] := 0.1466748;
   Prof_PriceDA.Data[3261] := 0.1466748;
   Prof_PriceDA.Data[3262] := 0.1466748;
   Prof_PriceDA.Data[3263] := 0.1466748;
   Prof_PriceDA.Data[3264] := 0.142992;
   Prof_PriceDA.Data[3265] := 0.142992;
   Prof_PriceDA.Data[3266] := 0.142992;
   Prof_PriceDA.Data[3267] := 0.142992;
   Prof_PriceDA.Data[3268] := 0.1355832;
   Prof_PriceDA.Data[3269] := 0.1355832;
   Prof_PriceDA.Data[3270] := 0.1355832;
   Prof_PriceDA.Data[3271] := 0.1355832;
   Prof_PriceDA.Data[3272] := 0.1330344;
   Prof_PriceDA.Data[3273] := 0.1330344;
   Prof_PriceDA.Data[3274] := 0.1330344;
   Prof_PriceDA.Data[3275] := 0.1330344;
   Prof_PriceDA.Data[3276] := 0.1339092;
   Prof_PriceDA.Data[3277] := 0.1339092;
   Prof_PriceDA.Data[3278] := 0.1339092;
   Prof_PriceDA.Data[3279] := 0.1339092;
   Prof_PriceDA.Data[3280] := 0.13311;
   Prof_PriceDA.Data[3281] := 0.13311;
   Prof_PriceDA.Data[3282] := 0.13311;
   Prof_PriceDA.Data[3283] := 0.13311;
   Prof_PriceDA.Data[3284] := 0.1378404;
   Prof_PriceDA.Data[3285] := 0.1378404;
   Prof_PriceDA.Data[3286] := 0.1378404;
   Prof_PriceDA.Data[3287] := 0.1378404;
   Prof_PriceDA.Data[3288] := 0.1674432;
   Prof_PriceDA.Data[3289] := 0.1674432;
   Prof_PriceDA.Data[3290] := 0.1674432;
   Prof_PriceDA.Data[3291] := 0.1674432;
   Prof_PriceDA.Data[3292] := 0.2056644;
   Prof_PriceDA.Data[3293] := 0.2056644;
   Prof_PriceDA.Data[3294] := 0.2056644;
   Prof_PriceDA.Data[3295] := 0.2056644;
   Prof_PriceDA.Data[3296] := 0.2289492;
   Prof_PriceDA.Data[3297] := 0.2289492;
   Prof_PriceDA.Data[3298] := 0.2289492;
   Prof_PriceDA.Data[3299] := 0.2289492;
   Prof_PriceDA.Data[3300] := 0.1763748;
   Prof_PriceDA.Data[3301] := 0.1763748;
   Prof_PriceDA.Data[3302] := 0.1763748;
   Prof_PriceDA.Data[3303] := 0.1763748;
   Prof_PriceDA.Data[3304] := 0.1474524;
   Prof_PriceDA.Data[3305] := 0.1474524;
   Prof_PriceDA.Data[3306] := 0.1474524;
   Prof_PriceDA.Data[3307] := 0.1474524;
   Prof_PriceDA.Data[3308] := 0.1369656;
   Prof_PriceDA.Data[3309] := 0.1369656;
   Prof_PriceDA.Data[3310] := 0.1369656;
   Prof_PriceDA.Data[3311] := 0.1369656;
   Prof_PriceDA.Data[3312] := 0.127602;
   Prof_PriceDA.Data[3313] := 0.127602;
   Prof_PriceDA.Data[3314] := 0.127602;
   Prof_PriceDA.Data[3315] := 0.127602;
   Prof_PriceDA.Data[3316] := 0.1222452;
   Prof_PriceDA.Data[3317] := 0.1222452;
   Prof_PriceDA.Data[3318] := 0.1222452;
   Prof_PriceDA.Data[3319] := 0.1222452;
   Prof_PriceDA.Data[3320] := 0.1296972;
   Prof_PriceDA.Data[3321] := 0.1296972;
   Prof_PriceDA.Data[3322] := 0.1296972;
   Prof_PriceDA.Data[3323] := 0.1296972;
   Prof_PriceDA.Data[3324] := 0.1542456;
   Prof_PriceDA.Data[3325] := 0.1542456;
   Prof_PriceDA.Data[3326] := 0.1542456;
   Prof_PriceDA.Data[3327] := 0.1542456;
   Prof_PriceDA.Data[3328] := 0.181332;
   Prof_PriceDA.Data[3329] := 0.181332;
   Prof_PriceDA.Data[3330] := 0.181332;
   Prof_PriceDA.Data[3331] := 0.181332;
   Prof_PriceDA.Data[3332] := 0.189324;
   Prof_PriceDA.Data[3333] := 0.189324;
   Prof_PriceDA.Data[3334] := 0.189324;
   Prof_PriceDA.Data[3335] := 0.189324;
   Prof_PriceDA.Data[3336] := 0.189;
   Prof_PriceDA.Data[3337] := 0.189;
   Prof_PriceDA.Data[3338] := 0.189;
   Prof_PriceDA.Data[3339] := 0.189;
   Prof_PriceDA.Data[3340] := 0.1863648;
   Prof_PriceDA.Data[3341] := 0.1863648;
   Prof_PriceDA.Data[3342] := 0.1863648;
   Prof_PriceDA.Data[3343] := 0.1863648;
   Prof_PriceDA.Data[3344] := 0.1727352;
   Prof_PriceDA.Data[3345] := 0.1727352;
   Prof_PriceDA.Data[3346] := 0.1727352;
   Prof_PriceDA.Data[3347] := 0.1727352;
   Prof_PriceDA.Data[3348] := 0.1464804;
   Prof_PriceDA.Data[3349] := 0.1464804;
   Prof_PriceDA.Data[3350] := 0.1464804;
   Prof_PriceDA.Data[3351] := 0.1464804;
   Prof_PriceDA.Data[3352] := 0.1424412;
   Prof_PriceDA.Data[3353] := 0.1424412;
   Prof_PriceDA.Data[3354] := 0.1424412;
   Prof_PriceDA.Data[3355] := 0.1424412;
   Prof_PriceDA.Data[3356] := 0.1347624;
   Prof_PriceDA.Data[3357] := 0.1347624;
   Prof_PriceDA.Data[3358] := 0.1347624;
   Prof_PriceDA.Data[3359] := 0.1347624;
   Prof_PriceDA.Data[3360] := 0.1260036;
   Prof_PriceDA.Data[3361] := 0.1260036;
   Prof_PriceDA.Data[3362] := 0.1260036;
   Prof_PriceDA.Data[3363] := 0.1260036;
   Prof_PriceDA.Data[3364] := 0.1207548;
   Prof_PriceDA.Data[3365] := 0.1207548;
   Prof_PriceDA.Data[3366] := 0.1207548;
   Prof_PriceDA.Data[3367] := 0.1207548;
   Prof_PriceDA.Data[3368] := 0.1198584;
   Prof_PriceDA.Data[3369] := 0.1198584;
   Prof_PriceDA.Data[3370] := 0.1198584;
   Prof_PriceDA.Data[3371] := 0.1198584;
   Prof_PriceDA.Data[3372] := 0.1186056;
   Prof_PriceDA.Data[3373] := 0.1186056;
   Prof_PriceDA.Data[3374] := 0.1186056;
   Prof_PriceDA.Data[3375] := 0.1186056;
   Prof_PriceDA.Data[3376] := 0.1248912;
   Prof_PriceDA.Data[3377] := 0.1248912;
   Prof_PriceDA.Data[3378] := 0.1248912;
   Prof_PriceDA.Data[3379] := 0.1248912;
   Prof_PriceDA.Data[3380] := 0.1323648;
   Prof_PriceDA.Data[3381] := 0.1323648;
   Prof_PriceDA.Data[3382] := 0.1323648;
   Prof_PriceDA.Data[3383] := 0.1323648;
   Prof_PriceDA.Data[3384] := 0.1636524;
   Prof_PriceDA.Data[3385] := 0.1636524;
   Prof_PriceDA.Data[3386] := 0.1636524;
   Prof_PriceDA.Data[3387] := 0.1636524;
   Prof_PriceDA.Data[3388] := 0.1825092;
   Prof_PriceDA.Data[3389] := 0.1825092;
   Prof_PriceDA.Data[3390] := 0.1825092;
   Prof_PriceDA.Data[3391] := 0.1825092;
   Prof_PriceDA.Data[3392] := 0.1952748;
   Prof_PriceDA.Data[3393] := 0.1952748;
   Prof_PriceDA.Data[3394] := 0.1952748;
   Prof_PriceDA.Data[3395] := 0.1952748;
   Prof_PriceDA.Data[3396] := 0.1720764;
   Prof_PriceDA.Data[3397] := 0.1720764;
   Prof_PriceDA.Data[3398] := 0.1720764;
   Prof_PriceDA.Data[3399] := 0.1720764;
   Prof_PriceDA.Data[3400] := 0.145476;
   Prof_PriceDA.Data[3401] := 0.145476;
   Prof_PriceDA.Data[3402] := 0.145476;
   Prof_PriceDA.Data[3403] := 0.145476;
   Prof_PriceDA.Data[3404] := 0.133704;
   Prof_PriceDA.Data[3405] := 0.133704;
   Prof_PriceDA.Data[3406] := 0.133704;
   Prof_PriceDA.Data[3407] := 0.133704;
   Prof_PriceDA.Data[3408] := 0.127926;
   Prof_PriceDA.Data[3409] := 0.127926;
   Prof_PriceDA.Data[3410] := 0.127926;
   Prof_PriceDA.Data[3411] := 0.127926;
   Prof_PriceDA.Data[3412] := 0.1297512;
   Prof_PriceDA.Data[3413] := 0.1297512;
   Prof_PriceDA.Data[3414] := 0.1297512;
   Prof_PriceDA.Data[3415] := 0.1297512;
   Prof_PriceDA.Data[3416] := 0.139158;
   Prof_PriceDA.Data[3417] := 0.139158;
   Prof_PriceDA.Data[3418] := 0.139158;
   Prof_PriceDA.Data[3419] := 0.139158;
   Prof_PriceDA.Data[3420] := 0.1556496;
   Prof_PriceDA.Data[3421] := 0.1556496;
   Prof_PriceDA.Data[3422] := 0.1556496;
   Prof_PriceDA.Data[3423] := 0.1556496;
   Prof_PriceDA.Data[3424] := 0.1719252;
   Prof_PriceDA.Data[3425] := 0.1719252;
   Prof_PriceDA.Data[3426] := 0.1719252;
   Prof_PriceDA.Data[3427] := 0.1719252;
   Prof_PriceDA.Data[3428] := 0.19116;
   Prof_PriceDA.Data[3429] := 0.19116;
   Prof_PriceDA.Data[3430] := 0.19116;
   Prof_PriceDA.Data[3431] := 0.19116;
   Prof_PriceDA.Data[3432] := 0.205092;
   Prof_PriceDA.Data[3433] := 0.205092;
   Prof_PriceDA.Data[3434] := 0.205092;
   Prof_PriceDA.Data[3435] := 0.205092;
   Prof_PriceDA.Data[3436] := 0.2048004;
   Prof_PriceDA.Data[3437] := 0.2048004;
   Prof_PriceDA.Data[3438] := 0.2048004;
   Prof_PriceDA.Data[3439] := 0.2048004;
   Prof_PriceDA.Data[3440] := 0.1836;
   Prof_PriceDA.Data[3441] := 0.1836;
   Prof_PriceDA.Data[3442] := 0.1836;
   Prof_PriceDA.Data[3443] := 0.1836;
   Prof_PriceDA.Data[3444] := 0.1678536;
   Prof_PriceDA.Data[3445] := 0.1678536;
   Prof_PriceDA.Data[3446] := 0.1678536;
   Prof_PriceDA.Data[3447] := 0.1678536;
   Prof_PriceDA.Data[3448] := 0.155196;
   Prof_PriceDA.Data[3449] := 0.155196;
   Prof_PriceDA.Data[3450] := 0.155196;
   Prof_PriceDA.Data[3451] := 0.155196;
   Prof_PriceDA.Data[3452] := 0.144774;
   Prof_PriceDA.Data[3453] := 0.144774;
   Prof_PriceDA.Data[3454] := 0.144774;
   Prof_PriceDA.Data[3455] := 0.144774;
   Prof_PriceDA.Data[3456] := 0.1443636;
   Prof_PriceDA.Data[3457] := 0.1443636;
   Prof_PriceDA.Data[3458] := 0.1443636;
   Prof_PriceDA.Data[3459] := 0.1443636;
   Prof_PriceDA.Data[3460] := 0.1403892;
   Prof_PriceDA.Data[3461] := 0.1403892;
   Prof_PriceDA.Data[3462] := 0.1403892;
   Prof_PriceDA.Data[3463] := 0.1403892;
   Prof_PriceDA.Data[3464] := 0.13608;
   Prof_PriceDA.Data[3465] := 0.13608;
   Prof_PriceDA.Data[3466] := 0.13608;
   Prof_PriceDA.Data[3467] := 0.13608;
   Prof_PriceDA.Data[3468] := 0.135;
   Prof_PriceDA.Data[3469] := 0.135;
   Prof_PriceDA.Data[3470] := 0.135;
   Prof_PriceDA.Data[3471] := 0.135;
   Prof_PriceDA.Data[3472] := 0.1350108;
   Prof_PriceDA.Data[3473] := 0.1350108;
   Prof_PriceDA.Data[3474] := 0.1350108;
   Prof_PriceDA.Data[3475] := 0.1350108;
   Prof_PriceDA.Data[3476] := 0.1447524;
   Prof_PriceDA.Data[3477] := 0.1447524;
   Prof_PriceDA.Data[3478] := 0.1447524;
   Prof_PriceDA.Data[3479] := 0.1447524;
   Prof_PriceDA.Data[3480] := 0.165996;
   Prof_PriceDA.Data[3481] := 0.165996;
   Prof_PriceDA.Data[3482] := 0.165996;
   Prof_PriceDA.Data[3483] := 0.165996;
   Prof_PriceDA.Data[3484] := 0.1944972;
   Prof_PriceDA.Data[3485] := 0.1944972;
   Prof_PriceDA.Data[3486] := 0.1944972;
   Prof_PriceDA.Data[3487] := 0.1944972;
   Prof_PriceDA.Data[3488] := 0.2356128;
   Prof_PriceDA.Data[3489] := 0.2356128;
   Prof_PriceDA.Data[3490] := 0.2356128;
   Prof_PriceDA.Data[3491] := 0.2356128;
   Prof_PriceDA.Data[3492] := 0.1930932;
   Prof_PriceDA.Data[3493] := 0.1930932;
   Prof_PriceDA.Data[3494] := 0.1930932;
   Prof_PriceDA.Data[3495] := 0.1930932;
   Prof_PriceDA.Data[3496] := 0.1686204;
   Prof_PriceDA.Data[3497] := 0.1686204;
   Prof_PriceDA.Data[3498] := 0.1686204;
   Prof_PriceDA.Data[3499] := 0.1686204;
   Prof_PriceDA.Data[3500] := 0.1617408;
   Prof_PriceDA.Data[3501] := 0.1617408;
   Prof_PriceDA.Data[3502] := 0.1617408;
   Prof_PriceDA.Data[3503] := 0.1617408;
   Prof_PriceDA.Data[3504] := 0.1561032;
   Prof_PriceDA.Data[3505] := 0.1561032;
   Prof_PriceDA.Data[3506] := 0.1561032;
   Prof_PriceDA.Data[3507] := 0.1561032;
   Prof_PriceDA.Data[3508] := 0.1526148;
   Prof_PriceDA.Data[3509] := 0.1526148;
   Prof_PriceDA.Data[3510] := 0.1526148;
   Prof_PriceDA.Data[3511] := 0.1526148;
   Prof_PriceDA.Data[3512] := 0.1520208;
   Prof_PriceDA.Data[3513] := 0.1520208;
   Prof_PriceDA.Data[3514] := 0.1520208;
   Prof_PriceDA.Data[3515] := 0.1520208;
   Prof_PriceDA.Data[3516] := 0.1622808;
   Prof_PriceDA.Data[3517] := 0.1622808;
   Prof_PriceDA.Data[3518] := 0.1622808;
   Prof_PriceDA.Data[3519] := 0.1622808;
   Prof_PriceDA.Data[3520] := 0.181656;
   Prof_PriceDA.Data[3521] := 0.181656;
   Prof_PriceDA.Data[3522] := 0.181656;
   Prof_PriceDA.Data[3523] := 0.181656;
   Prof_PriceDA.Data[3524] := 0.188244;
   Prof_PriceDA.Data[3525] := 0.188244;
   Prof_PriceDA.Data[3526] := 0.188244;
   Prof_PriceDA.Data[3527] := 0.188244;
   Prof_PriceDA.Data[3528] := 0.1913544;
   Prof_PriceDA.Data[3529] := 0.1913544;
   Prof_PriceDA.Data[3530] := 0.1913544;
   Prof_PriceDA.Data[3531] := 0.1913544;
   Prof_PriceDA.Data[3532] := 0.1864512;
   Prof_PriceDA.Data[3533] := 0.1864512;
   Prof_PriceDA.Data[3534] := 0.1864512;
   Prof_PriceDA.Data[3535] := 0.1864512;
   Prof_PriceDA.Data[3536] := 0.1768068;
   Prof_PriceDA.Data[3537] := 0.1768068;
   Prof_PriceDA.Data[3538] := 0.1768068;
   Prof_PriceDA.Data[3539] := 0.1768068;
   Prof_PriceDA.Data[3540] := 0.159624;
   Prof_PriceDA.Data[3541] := 0.159624;
   Prof_PriceDA.Data[3542] := 0.159624;
   Prof_PriceDA.Data[3543] := 0.159624;
   Prof_PriceDA.Data[3544] := 0.1512108;
   Prof_PriceDA.Data[3545] := 0.1512108;
   Prof_PriceDA.Data[3546] := 0.1512108;
   Prof_PriceDA.Data[3547] := 0.1512108;
   Prof_PriceDA.Data[3548] := 0.131706;
   Prof_PriceDA.Data[3549] := 0.131706;
   Prof_PriceDA.Data[3550] := 0.131706;
   Prof_PriceDA.Data[3551] := 0.131706;
   Prof_PriceDA.Data[3552] := 0.136134;
   Prof_PriceDA.Data[3553] := 0.136134;
   Prof_PriceDA.Data[3554] := 0.136134;
   Prof_PriceDA.Data[3555] := 0.136134;
   Prof_PriceDA.Data[3556] := 0.121716;
   Prof_PriceDA.Data[3557] := 0.121716;
   Prof_PriceDA.Data[3558] := 0.121716;
   Prof_PriceDA.Data[3559] := 0.121716;
   Prof_PriceDA.Data[3560] := 0.1175256;
   Prof_PriceDA.Data[3561] := 0.1175256;
   Prof_PriceDA.Data[3562] := 0.1175256;
   Prof_PriceDA.Data[3563] := 0.1175256;
   Prof_PriceDA.Data[3564] := 0.1134;
   Prof_PriceDA.Data[3565] := 0.1134;
   Prof_PriceDA.Data[3566] := 0.1134;
   Prof_PriceDA.Data[3567] := 0.1134;
   Prof_PriceDA.Data[3568] := 0.1185192;
   Prof_PriceDA.Data[3569] := 0.1185192;
   Prof_PriceDA.Data[3570] := 0.1185192;
   Prof_PriceDA.Data[3571] := 0.1185192;
   Prof_PriceDA.Data[3572] := 0.1280772;
   Prof_PriceDA.Data[3573] := 0.1280772;
   Prof_PriceDA.Data[3574] := 0.1280772;
   Prof_PriceDA.Data[3575] := 0.1280772;
   Prof_PriceDA.Data[3576] := 0.1678104;
   Prof_PriceDA.Data[3577] := 0.1678104;
   Prof_PriceDA.Data[3578] := 0.1678104;
   Prof_PriceDA.Data[3579] := 0.1678104;
   Prof_PriceDA.Data[3580] := 0.1848744;
   Prof_PriceDA.Data[3581] := 0.1848744;
   Prof_PriceDA.Data[3582] := 0.1848744;
   Prof_PriceDA.Data[3583] := 0.1848744;
   Prof_PriceDA.Data[3584] := 0.1782324;
   Prof_PriceDA.Data[3585] := 0.1782324;
   Prof_PriceDA.Data[3586] := 0.1782324;
   Prof_PriceDA.Data[3587] := 0.1782324;
   Prof_PriceDA.Data[3588] := 0.1625076;
   Prof_PriceDA.Data[3589] := 0.1625076;
   Prof_PriceDA.Data[3590] := 0.1625076;
   Prof_PriceDA.Data[3591] := 0.1625076;
   Prof_PriceDA.Data[3592] := 0.1456812;
   Prof_PriceDA.Data[3593] := 0.1456812;
   Prof_PriceDA.Data[3594] := 0.1456812;
   Prof_PriceDA.Data[3595] := 0.1456812;
   Prof_PriceDA.Data[3596] := 0.1280556;
   Prof_PriceDA.Data[3597] := 0.1280556;
   Prof_PriceDA.Data[3598] := 0.1280556;
   Prof_PriceDA.Data[3599] := 0.1280556;
   Prof_PriceDA.Data[3600] := 0.1243512;
   Prof_PriceDA.Data[3601] := 0.1243512;
   Prof_PriceDA.Data[3602] := 0.1243512;
   Prof_PriceDA.Data[3603] := 0.1243512;
   Prof_PriceDA.Data[3604] := 0.1240164;
   Prof_PriceDA.Data[3605] := 0.1240164;
   Prof_PriceDA.Data[3606] := 0.1240164;
   Prof_PriceDA.Data[3607] := 0.1240164;
   Prof_PriceDA.Data[3608] := 0.12744;
   Prof_PriceDA.Data[3609] := 0.12744;
   Prof_PriceDA.Data[3610] := 0.12744;
   Prof_PriceDA.Data[3611] := 0.12744;
   Prof_PriceDA.Data[3612] := 0.1442556;
   Prof_PriceDA.Data[3613] := 0.1442556;
   Prof_PriceDA.Data[3614] := 0.1442556;
   Prof_PriceDA.Data[3615] := 0.1442556;
   Prof_PriceDA.Data[3616] := 0.1857924;
   Prof_PriceDA.Data[3617] := 0.1857924;
   Prof_PriceDA.Data[3618] := 0.1857924;
   Prof_PriceDA.Data[3619] := 0.1857924;
   Prof_PriceDA.Data[3620] := 0.1894644;
   Prof_PriceDA.Data[3621] := 0.1894644;
   Prof_PriceDA.Data[3622] := 0.1894644;
   Prof_PriceDA.Data[3623] := 0.1894644;
   Prof_PriceDA.Data[3624] := 0.1884924;
   Prof_PriceDA.Data[3625] := 0.1884924;
   Prof_PriceDA.Data[3626] := 0.1884924;
   Prof_PriceDA.Data[3627] := 0.1884924;
   Prof_PriceDA.Data[3628] := 0.1860624;
   Prof_PriceDA.Data[3629] := 0.1860624;
   Prof_PriceDA.Data[3630] := 0.1860624;
   Prof_PriceDA.Data[3631] := 0.1860624;
   Prof_PriceDA.Data[3632] := 0.1818072;
   Prof_PriceDA.Data[3633] := 0.1818072;
   Prof_PriceDA.Data[3634] := 0.1818072;
   Prof_PriceDA.Data[3635] := 0.1818072;
   Prof_PriceDA.Data[3636] := 0.1557576;
   Prof_PriceDA.Data[3637] := 0.1557576;
   Prof_PriceDA.Data[3638] := 0.1557576;
   Prof_PriceDA.Data[3639] := 0.1557576;
   Prof_PriceDA.Data[3640] := 0.1285632;
   Prof_PriceDA.Data[3641] := 0.1285632;
   Prof_PriceDA.Data[3642] := 0.1285632;
   Prof_PriceDA.Data[3643] := 0.1285632;
   Prof_PriceDA.Data[3644] := 0.1209816;
   Prof_PriceDA.Data[3645] := 0.1209816;
   Prof_PriceDA.Data[3646] := 0.1209816;
   Prof_PriceDA.Data[3647] := 0.1209816;
   Prof_PriceDA.Data[3648] := 0.09828;
   Prof_PriceDA.Data[3649] := 0.09828;
   Prof_PriceDA.Data[3650] := 0.09828;
   Prof_PriceDA.Data[3651] := 0.09828;
   Prof_PriceDA.Data[3652] := 0.0950184;
   Prof_PriceDA.Data[3653] := 0.0950184;
   Prof_PriceDA.Data[3654] := 0.0950184;
   Prof_PriceDA.Data[3655] := 0.0950184;
   Prof_PriceDA.Data[3656] := 0.0937872;
   Prof_PriceDA.Data[3657] := 0.0937872;
   Prof_PriceDA.Data[3658] := 0.0937872;
   Prof_PriceDA.Data[3659] := 0.0937872;
   Prof_PriceDA.Data[3660] := 0.09612;
   Prof_PriceDA.Data[3661] := 0.09612;
   Prof_PriceDA.Data[3662] := 0.09612;
   Prof_PriceDA.Data[3663] := 0.09612;
   Prof_PriceDA.Data[3664] := 0.0968652;
   Prof_PriceDA.Data[3665] := 0.0968652;
   Prof_PriceDA.Data[3666] := 0.0968652;
   Prof_PriceDA.Data[3667] := 0.0968652;
   Prof_PriceDA.Data[3668] := 0.0982692;
   Prof_PriceDA.Data[3669] := 0.0982692;
   Prof_PriceDA.Data[3670] := 0.0982692;
   Prof_PriceDA.Data[3671] := 0.0982692;
   Prof_PriceDA.Data[3672] := 0.1052028;
   Prof_PriceDA.Data[3673] := 0.1052028;
   Prof_PriceDA.Data[3674] := 0.1052028;
   Prof_PriceDA.Data[3675] := 0.1052028;
   Prof_PriceDA.Data[3676] := 0.1174068;
   Prof_PriceDA.Data[3677] := 0.1174068;
   Prof_PriceDA.Data[3678] := 0.1174068;
   Prof_PriceDA.Data[3679] := 0.1174068;
   Prof_PriceDA.Data[3680] := 0.1222128;
   Prof_PriceDA.Data[3681] := 0.1222128;
   Prof_PriceDA.Data[3682] := 0.1222128;
   Prof_PriceDA.Data[3683] := 0.1222128;
   Prof_PriceDA.Data[3684] := 0.109134;
   Prof_PriceDA.Data[3685] := 0.109134;
   Prof_PriceDA.Data[3686] := 0.109134;
   Prof_PriceDA.Data[3687] := 0.109134;
   Prof_PriceDA.Data[3688] := 0.1035072;
   Prof_PriceDA.Data[3689] := 0.1035072;
   Prof_PriceDA.Data[3690] := 0.1035072;
   Prof_PriceDA.Data[3691] := 0.1035072;
   Prof_PriceDA.Data[3692] := 0.0960336;
   Prof_PriceDA.Data[3693] := 0.0960336;
   Prof_PriceDA.Data[3694] := 0.0960336;
   Prof_PriceDA.Data[3695] := 0.0960336;
   Prof_PriceDA.Data[3696] := 0.0954828;
   Prof_PriceDA.Data[3697] := 0.0954828;
   Prof_PriceDA.Data[3698] := 0.0954828;
   Prof_PriceDA.Data[3699] := 0.0954828;
   Prof_PriceDA.Data[3700] := 0.097686;
   Prof_PriceDA.Data[3701] := 0.097686;
   Prof_PriceDA.Data[3702] := 0.097686;
   Prof_PriceDA.Data[3703] := 0.097686;
   Prof_PriceDA.Data[3704] := 0.1025244;
   Prof_PriceDA.Data[3705] := 0.1025244;
   Prof_PriceDA.Data[3706] := 0.1025244;
   Prof_PriceDA.Data[3707] := 0.1025244;
   Prof_PriceDA.Data[3708] := 0.12744;
   Prof_PriceDA.Data[3709] := 0.12744;
   Prof_PriceDA.Data[3710] := 0.12744;
   Prof_PriceDA.Data[3711] := 0.12744;
   Prof_PriceDA.Data[3712] := 0.16173;
   Prof_PriceDA.Data[3713] := 0.16173;
   Prof_PriceDA.Data[3714] := 0.16173;
   Prof_PriceDA.Data[3715] := 0.16173;
   Prof_PriceDA.Data[3716] := 0.1752948;
   Prof_PriceDA.Data[3717] := 0.1752948;
   Prof_PriceDA.Data[3718] := 0.1752948;
   Prof_PriceDA.Data[3719] := 0.1752948;
   Prof_PriceDA.Data[3720] := 0.1733832;
   Prof_PriceDA.Data[3721] := 0.1733832;
   Prof_PriceDA.Data[3722] := 0.1733832;
   Prof_PriceDA.Data[3723] := 0.1733832;
   Prof_PriceDA.Data[3724] := 0.1713852;
   Prof_PriceDA.Data[3725] := 0.1713852;
   Prof_PriceDA.Data[3726] := 0.1713852;
   Prof_PriceDA.Data[3727] := 0.1713852;
   Prof_PriceDA.Data[3728] := 0.1661472;
   Prof_PriceDA.Data[3729] := 0.1661472;
   Prof_PriceDA.Data[3730] := 0.1661472;
   Prof_PriceDA.Data[3731] := 0.1661472;
   Prof_PriceDA.Data[3732] := 0.16092;
   Prof_PriceDA.Data[3733] := 0.16092;
   Prof_PriceDA.Data[3734] := 0.16092;
   Prof_PriceDA.Data[3735] := 0.16092;
   Prof_PriceDA.Data[3736] := 0.1542564;
   Prof_PriceDA.Data[3737] := 0.1542564;
   Prof_PriceDA.Data[3738] := 0.1542564;
   Prof_PriceDA.Data[3739] := 0.1542564;
   Prof_PriceDA.Data[3740] := 0.1449792;
   Prof_PriceDA.Data[3741] := 0.1449792;
   Prof_PriceDA.Data[3742] := 0.1449792;
   Prof_PriceDA.Data[3743] := 0.1449792;
   Prof_PriceDA.Data[3744] := 0.1458;
   Prof_PriceDA.Data[3745] := 0.1458;
   Prof_PriceDA.Data[3746] := 0.1458;
   Prof_PriceDA.Data[3747] := 0.1458;
   Prof_PriceDA.Data[3748] := 0.136404;
   Prof_PriceDA.Data[3749] := 0.136404;
   Prof_PriceDA.Data[3750] := 0.136404;
   Prof_PriceDA.Data[3751] := 0.136404;
   Prof_PriceDA.Data[3752] := 0.1319004;
   Prof_PriceDA.Data[3753] := 0.1319004;
   Prof_PriceDA.Data[3754] := 0.1319004;
   Prof_PriceDA.Data[3755] := 0.1319004;
   Prof_PriceDA.Data[3756] := 0.128844;
   Prof_PriceDA.Data[3757] := 0.128844;
   Prof_PriceDA.Data[3758] := 0.128844;
   Prof_PriceDA.Data[3759] := 0.128844;
   Prof_PriceDA.Data[3760] := 0.1261656;
   Prof_PriceDA.Data[3761] := 0.1261656;
   Prof_PriceDA.Data[3762] := 0.1261656;
   Prof_PriceDA.Data[3763] := 0.1261656;
   Prof_PriceDA.Data[3764] := 0.12636;
   Prof_PriceDA.Data[3765] := 0.12636;
   Prof_PriceDA.Data[3766] := 0.12636;
   Prof_PriceDA.Data[3767] := 0.12636;
   Prof_PriceDA.Data[3768] := 0.12636;
   Prof_PriceDA.Data[3769] := 0.12636;
   Prof_PriceDA.Data[3770] := 0.12636;
   Prof_PriceDA.Data[3771] := 0.12636;
   Prof_PriceDA.Data[3772] := 0.1441044;
   Prof_PriceDA.Data[3773] := 0.1441044;
   Prof_PriceDA.Data[3774] := 0.1441044;
   Prof_PriceDA.Data[3775] := 0.1441044;
   Prof_PriceDA.Data[3776] := 0.1477116;
   Prof_PriceDA.Data[3777] := 0.1477116;
   Prof_PriceDA.Data[3778] := 0.1477116;
   Prof_PriceDA.Data[3779] := 0.1477116;
   Prof_PriceDA.Data[3780] := 0.1321812;
   Prof_PriceDA.Data[3781] := 0.1321812;
   Prof_PriceDA.Data[3782] := 0.1321812;
   Prof_PriceDA.Data[3783] := 0.1321812;
   Prof_PriceDA.Data[3784] := 0.1230876;
   Prof_PriceDA.Data[3785] := 0.1230876;
   Prof_PriceDA.Data[3786] := 0.1230876;
   Prof_PriceDA.Data[3787] := 0.1230876;
   Prof_PriceDA.Data[3788] := 0.1191456;
   Prof_PriceDA.Data[3789] := 0.1191456;
   Prof_PriceDA.Data[3790] := 0.1191456;
   Prof_PriceDA.Data[3791] := 0.1191456;
   Prof_PriceDA.Data[3792] := 0.1106028;
   Prof_PriceDA.Data[3793] := 0.1106028;
   Prof_PriceDA.Data[3794] := 0.1106028;
   Prof_PriceDA.Data[3795] := 0.1106028;
   Prof_PriceDA.Data[3796] := 0.1090368;
   Prof_PriceDA.Data[3797] := 0.1090368;
   Prof_PriceDA.Data[3798] := 0.1090368;
   Prof_PriceDA.Data[3799] := 0.1090368;
   Prof_PriceDA.Data[3800] := 0.118692;
   Prof_PriceDA.Data[3801] := 0.118692;
   Prof_PriceDA.Data[3802] := 0.118692;
   Prof_PriceDA.Data[3803] := 0.118692;
   Prof_PriceDA.Data[3804] := 0.130032;
   Prof_PriceDA.Data[3805] := 0.130032;
   Prof_PriceDA.Data[3806] := 0.130032;
   Prof_PriceDA.Data[3807] := 0.130032;
   Prof_PriceDA.Data[3808] := 0.1627992;
   Prof_PriceDA.Data[3809] := 0.1627992;
   Prof_PriceDA.Data[3810] := 0.1627992;
   Prof_PriceDA.Data[3811] := 0.1627992;
   Prof_PriceDA.Data[3812] := 0.1736856;
   Prof_PriceDA.Data[3813] := 0.1736856;
   Prof_PriceDA.Data[3814] := 0.1736856;
   Prof_PriceDA.Data[3815] := 0.1736856;
   Prof_PriceDA.Data[3816] := 0.1889784;
   Prof_PriceDA.Data[3817] := 0.1889784;
   Prof_PriceDA.Data[3818] := 0.1889784;
   Prof_PriceDA.Data[3819] := 0.1889784;
   Prof_PriceDA.Data[3820] := 0.1888164;
   Prof_PriceDA.Data[3821] := 0.1888164;
   Prof_PriceDA.Data[3822] := 0.1888164;
   Prof_PriceDA.Data[3823] := 0.1888164;
   Prof_PriceDA.Data[3824] := 0.1786968;
   Prof_PriceDA.Data[3825] := 0.1786968;
   Prof_PriceDA.Data[3826] := 0.1786968;
   Prof_PriceDA.Data[3827] := 0.1786968;
   Prof_PriceDA.Data[3828] := 0.1560816;
   Prof_PriceDA.Data[3829] := 0.1560816;
   Prof_PriceDA.Data[3830] := 0.1560816;
   Prof_PriceDA.Data[3831] := 0.1560816;
   Prof_PriceDA.Data[3832] := 0.15444;
   Prof_PriceDA.Data[3833] := 0.15444;
   Prof_PriceDA.Data[3834] := 0.15444;
   Prof_PriceDA.Data[3835] := 0.15444;
   Prof_PriceDA.Data[3836] := 0.139482;
   Prof_PriceDA.Data[3837] := 0.139482;
   Prof_PriceDA.Data[3838] := 0.139482;
   Prof_PriceDA.Data[3839] := 0.139482;
   Prof_PriceDA.Data[3840] := 0.1297944;
   Prof_PriceDA.Data[3841] := 0.1297944;
   Prof_PriceDA.Data[3842] := 0.1297944;
   Prof_PriceDA.Data[3843] := 0.1297944;
   Prof_PriceDA.Data[3844] := 0.1247292;
   Prof_PriceDA.Data[3845] := 0.1247292;
   Prof_PriceDA.Data[3846] := 0.1247292;
   Prof_PriceDA.Data[3847] := 0.1247292;
   Prof_PriceDA.Data[3848] := 0.1217916;
   Prof_PriceDA.Data[3849] := 0.1217916;
   Prof_PriceDA.Data[3850] := 0.1217916;
   Prof_PriceDA.Data[3851] := 0.1217916;
   Prof_PriceDA.Data[3852] := 0.1173096;
   Prof_PriceDA.Data[3853] := 0.1173096;
   Prof_PriceDA.Data[3854] := 0.1173096;
   Prof_PriceDA.Data[3855] := 0.1173096;
   Prof_PriceDA.Data[3856] := 0.1168992;
   Prof_PriceDA.Data[3857] := 0.1168992;
   Prof_PriceDA.Data[3858] := 0.1168992;
   Prof_PriceDA.Data[3859] := 0.1168992;
   Prof_PriceDA.Data[3860] := 0.126576;
   Prof_PriceDA.Data[3861] := 0.126576;
   Prof_PriceDA.Data[3862] := 0.126576;
   Prof_PriceDA.Data[3863] := 0.126576;
   Prof_PriceDA.Data[3864] := 0.1724004;
   Prof_PriceDA.Data[3865] := 0.1724004;
   Prof_PriceDA.Data[3866] := 0.1724004;
   Prof_PriceDA.Data[3867] := 0.1724004;
   Prof_PriceDA.Data[3868] := 0.1935684;
   Prof_PriceDA.Data[3869] := 0.1935684;
   Prof_PriceDA.Data[3870] := 0.1935684;
   Prof_PriceDA.Data[3871] := 0.1935684;
   Prof_PriceDA.Data[3872] := 0.1958688;
   Prof_PriceDA.Data[3873] := 0.1958688;
   Prof_PriceDA.Data[3874] := 0.1958688;
   Prof_PriceDA.Data[3875] := 0.1958688;
   Prof_PriceDA.Data[3876] := 0.1762344;
   Prof_PriceDA.Data[3877] := 0.1762344;
   Prof_PriceDA.Data[3878] := 0.1762344;
   Prof_PriceDA.Data[3879] := 0.1762344;
   Prof_PriceDA.Data[3880] := 0.1672488;
   Prof_PriceDA.Data[3881] := 0.1672488;
   Prof_PriceDA.Data[3882] := 0.1672488;
   Prof_PriceDA.Data[3883] := 0.1672488;
   Prof_PriceDA.Data[3884] := 0.1512108;
   Prof_PriceDA.Data[3885] := 0.1512108;
   Prof_PriceDA.Data[3886] := 0.1512108;
   Prof_PriceDA.Data[3887] := 0.1512108;
   Prof_PriceDA.Data[3888] := 0.136512;
   Prof_PriceDA.Data[3889] := 0.136512;
   Prof_PriceDA.Data[3890] := 0.136512;
   Prof_PriceDA.Data[3891] := 0.136512;
   Prof_PriceDA.Data[3892] := 0.132732;
   Prof_PriceDA.Data[3893] := 0.132732;
   Prof_PriceDA.Data[3894] := 0.132732;
   Prof_PriceDA.Data[3895] := 0.132732;
   Prof_PriceDA.Data[3896] := 0.142398;
   Prof_PriceDA.Data[3897] := 0.142398;
   Prof_PriceDA.Data[3898] := 0.142398;
   Prof_PriceDA.Data[3899] := 0.142398;
   Prof_PriceDA.Data[3900] := 0.179712;
   Prof_PriceDA.Data[3901] := 0.179712;
   Prof_PriceDA.Data[3902] := 0.179712;
   Prof_PriceDA.Data[3903] := 0.179712;
   Prof_PriceDA.Data[3904] := 0.2052972;
   Prof_PriceDA.Data[3905] := 0.2052972;
   Prof_PriceDA.Data[3906] := 0.2052972;
   Prof_PriceDA.Data[3907] := 0.2052972;
   Prof_PriceDA.Data[3908] := 0.218322;
   Prof_PriceDA.Data[3909] := 0.218322;
   Prof_PriceDA.Data[3910] := 0.218322;
   Prof_PriceDA.Data[3911] := 0.218322;
   Prof_PriceDA.Data[3912] := 0.2210112;
   Prof_PriceDA.Data[3913] := 0.2210112;
   Prof_PriceDA.Data[3914] := 0.2210112;
   Prof_PriceDA.Data[3915] := 0.2210112;
   Prof_PriceDA.Data[3916] := 0.2083752;
   Prof_PriceDA.Data[3917] := 0.2083752;
   Prof_PriceDA.Data[3918] := 0.2083752;
   Prof_PriceDA.Data[3919] := 0.2083752;
   Prof_PriceDA.Data[3920] := 0.2056644;
   Prof_PriceDA.Data[3921] := 0.2056644;
   Prof_PriceDA.Data[3922] := 0.2056644;
   Prof_PriceDA.Data[3923] := 0.2056644;
   Prof_PriceDA.Data[3924] := 0.1809;
   Prof_PriceDA.Data[3925] := 0.1809;
   Prof_PriceDA.Data[3926] := 0.1809;
   Prof_PriceDA.Data[3927] := 0.1809;
   Prof_PriceDA.Data[3928] := 0.1751544;
   Prof_PriceDA.Data[3929] := 0.1751544;
   Prof_PriceDA.Data[3930] := 0.1751544;
   Prof_PriceDA.Data[3931] := 0.1751544;
   Prof_PriceDA.Data[3932] := 0.1435428;
   Prof_PriceDA.Data[3933] := 0.1435428;
   Prof_PriceDA.Data[3934] := 0.1435428;
   Prof_PriceDA.Data[3935] := 0.1435428;
   Prof_PriceDA.Data[3936] := 0.1483812;
   Prof_PriceDA.Data[3937] := 0.1483812;
   Prof_PriceDA.Data[3938] := 0.1483812;
   Prof_PriceDA.Data[3939] := 0.1483812;
   Prof_PriceDA.Data[3940] := 0.1365768;
   Prof_PriceDA.Data[3941] := 0.1365768;
   Prof_PriceDA.Data[3942] := 0.1365768;
   Prof_PriceDA.Data[3943] := 0.1365768;
   Prof_PriceDA.Data[3944] := 0.1335204;
   Prof_PriceDA.Data[3945] := 0.1335204;
   Prof_PriceDA.Data[3946] := 0.1335204;
   Prof_PriceDA.Data[3947] := 0.1335204;
   Prof_PriceDA.Data[3948] := 0.1290384;
   Prof_PriceDA.Data[3949] := 0.1290384;
   Prof_PriceDA.Data[3950] := 0.1290384;
   Prof_PriceDA.Data[3951] := 0.1290384;
   Prof_PriceDA.Data[3952] := 0.1365876;
   Prof_PriceDA.Data[3953] := 0.1365876;
   Prof_PriceDA.Data[3954] := 0.1365876;
   Prof_PriceDA.Data[3955] := 0.1365876;
   Prof_PriceDA.Data[3956] := 0.1763856;
   Prof_PriceDA.Data[3957] := 0.1763856;
   Prof_PriceDA.Data[3958] := 0.1763856;
   Prof_PriceDA.Data[3959] := 0.1763856;
   Prof_PriceDA.Data[3960] := 0.1951884;
   Prof_PriceDA.Data[3961] := 0.1951884;
   Prof_PriceDA.Data[3962] := 0.1951884;
   Prof_PriceDA.Data[3963] := 0.1951884;
   Prof_PriceDA.Data[3964] := 0.2572236;
   Prof_PriceDA.Data[3965] := 0.2572236;
   Prof_PriceDA.Data[3966] := 0.2572236;
   Prof_PriceDA.Data[3967] := 0.2572236;
   Prof_PriceDA.Data[3968] := 0.1924884;
   Prof_PriceDA.Data[3969] := 0.1924884;
   Prof_PriceDA.Data[3970] := 0.1924884;
   Prof_PriceDA.Data[3971] := 0.1924884;
   Prof_PriceDA.Data[3972] := 0.15687;
   Prof_PriceDA.Data[3973] := 0.15687;
   Prof_PriceDA.Data[3974] := 0.15687;
   Prof_PriceDA.Data[3975] := 0.15687;
   Prof_PriceDA.Data[3976] := 0.13068;
   Prof_PriceDA.Data[3977] := 0.13068;
   Prof_PriceDA.Data[3978] := 0.13068;
   Prof_PriceDA.Data[3979] := 0.13068;
   Prof_PriceDA.Data[3980] := 0.1269432;
   Prof_PriceDA.Data[3981] := 0.1269432;
   Prof_PriceDA.Data[3982] := 0.1269432;
   Prof_PriceDA.Data[3983] := 0.1269432;
   Prof_PriceDA.Data[3984] := 0.1278612;
   Prof_PriceDA.Data[3985] := 0.1278612;
   Prof_PriceDA.Data[3986] := 0.1278612;
   Prof_PriceDA.Data[3987] := 0.1278612;
   Prof_PriceDA.Data[3988] := 0.1289304;
   Prof_PriceDA.Data[3989] := 0.1289304;
   Prof_PriceDA.Data[3990] := 0.1289304;
   Prof_PriceDA.Data[3991] := 0.1289304;
   Prof_PriceDA.Data[3992] := 0.1395684;
   Prof_PriceDA.Data[3993] := 0.1395684;
   Prof_PriceDA.Data[3994] := 0.1395684;
   Prof_PriceDA.Data[3995] := 0.1395684;
   Prof_PriceDA.Data[3996] := 0.1727136;
   Prof_PriceDA.Data[3997] := 0.1727136;
   Prof_PriceDA.Data[3998] := 0.1727136;
   Prof_PriceDA.Data[3999] := 0.1727136;
   Prof_PriceDA.Data[4000] := 0.200016;
   Prof_PriceDA.Data[4001] := 0.200016;
   Prof_PriceDA.Data[4002] := 0.200016;
   Prof_PriceDA.Data[4003] := 0.200016;
   Prof_PriceDA.Data[4004] := 0.2052;
   Prof_PriceDA.Data[4005] := 0.2052;
   Prof_PriceDA.Data[4006] := 0.2052;
   Prof_PriceDA.Data[4007] := 0.2052;
   Prof_PriceDA.Data[4008] := 0.2388312;
   Prof_PriceDA.Data[4009] := 0.2388312;
   Prof_PriceDA.Data[4010] := 0.2388312;
   Prof_PriceDA.Data[4011] := 0.2388312;
   Prof_PriceDA.Data[4012] := 0.2170044;
   Prof_PriceDA.Data[4013] := 0.2170044;
   Prof_PriceDA.Data[4014] := 0.2170044;
   Prof_PriceDA.Data[4015] := 0.2170044;
   Prof_PriceDA.Data[4016] := 0.1934064;
   Prof_PriceDA.Data[4017] := 0.1934064;
   Prof_PriceDA.Data[4018] := 0.1934064;
   Prof_PriceDA.Data[4019] := 0.1934064;
   Prof_PriceDA.Data[4020] := 0.1859868;
   Prof_PriceDA.Data[4021] := 0.1859868;
   Prof_PriceDA.Data[4022] := 0.1859868;
   Prof_PriceDA.Data[4023] := 0.1859868;
   Prof_PriceDA.Data[4024] := 0.1727892;
   Prof_PriceDA.Data[4025] := 0.1727892;
   Prof_PriceDA.Data[4026] := 0.1727892;
   Prof_PriceDA.Data[4027] := 0.1727892;
   Prof_PriceDA.Data[4028] := 0.1431432;
   Prof_PriceDA.Data[4029] := 0.1431432;
   Prof_PriceDA.Data[4030] := 0.1431432;
   Prof_PriceDA.Data[4031] := 0.1431432;
   Prof_PriceDA.Data[4032] := 0.1397952;
   Prof_PriceDA.Data[4033] := 0.1397952;
   Prof_PriceDA.Data[4034] := 0.1397952;
   Prof_PriceDA.Data[4035] := 0.1397952;
   Prof_PriceDA.Data[4036] := 0.1380996;
   Prof_PriceDA.Data[4037] := 0.1380996;
   Prof_PriceDA.Data[4038] := 0.1380996;
   Prof_PriceDA.Data[4039] := 0.1380996;
   Prof_PriceDA.Data[4040] := 0.1369656;
   Prof_PriceDA.Data[4041] := 0.1369656;
   Prof_PriceDA.Data[4042] := 0.1369656;
   Prof_PriceDA.Data[4043] := 0.1369656;
   Prof_PriceDA.Data[4044] := 0.1367172;
   Prof_PriceDA.Data[4045] := 0.1367172;
   Prof_PriceDA.Data[4046] := 0.1367172;
   Prof_PriceDA.Data[4047] := 0.1367172;
   Prof_PriceDA.Data[4048] := 0.1390392;
   Prof_PriceDA.Data[4049] := 0.1390392;
   Prof_PriceDA.Data[4050] := 0.1390392;
   Prof_PriceDA.Data[4051] := 0.1390392;
   Prof_PriceDA.Data[4052] := 0.1469772;
   Prof_PriceDA.Data[4053] := 0.1469772;
   Prof_PriceDA.Data[4054] := 0.1469772;
   Prof_PriceDA.Data[4055] := 0.1469772;
   Prof_PriceDA.Data[4056] := 0.1866024;
   Prof_PriceDA.Data[4057] := 0.1866024;
   Prof_PriceDA.Data[4058] := 0.1866024;
   Prof_PriceDA.Data[4059] := 0.1866024;
   Prof_PriceDA.Data[4060] := 0.1955232;
   Prof_PriceDA.Data[4061] := 0.1955232;
   Prof_PriceDA.Data[4062] := 0.1955232;
   Prof_PriceDA.Data[4063] := 0.1955232;
   Prof_PriceDA.Data[4064] := 0.1944;
   Prof_PriceDA.Data[4065] := 0.1944;
   Prof_PriceDA.Data[4066] := 0.1944;
   Prof_PriceDA.Data[4067] := 0.1944;
   Prof_PriceDA.Data[4068] := 0.1889136;
   Prof_PriceDA.Data[4069] := 0.1889136;
   Prof_PriceDA.Data[4070] := 0.1889136;
   Prof_PriceDA.Data[4071] := 0.1889136;
   Prof_PriceDA.Data[4072] := 0.1791612;
   Prof_PriceDA.Data[4073] := 0.1791612;
   Prof_PriceDA.Data[4074] := 0.1791612;
   Prof_PriceDA.Data[4075] := 0.1791612;
   Prof_PriceDA.Data[4076] := 0.171234;
   Prof_PriceDA.Data[4077] := 0.171234;
   Prof_PriceDA.Data[4078] := 0.171234;
   Prof_PriceDA.Data[4079] := 0.171234;
   Prof_PriceDA.Data[4080] := 0.16119;
   Prof_PriceDA.Data[4081] := 0.16119;
   Prof_PriceDA.Data[4082] := 0.16119;
   Prof_PriceDA.Data[4083] := 0.16119;
   Prof_PriceDA.Data[4084] := 0.1638144;
   Prof_PriceDA.Data[4085] := 0.1638144;
   Prof_PriceDA.Data[4086] := 0.1638144;
   Prof_PriceDA.Data[4087] := 0.1638144;
   Prof_PriceDA.Data[4088] := 0.1802196;
   Prof_PriceDA.Data[4089] := 0.1802196;
   Prof_PriceDA.Data[4090] := 0.1802196;
   Prof_PriceDA.Data[4091] := 0.1802196;
   Prof_PriceDA.Data[4092] := 0.1956852;
   Prof_PriceDA.Data[4093] := 0.1956852;
   Prof_PriceDA.Data[4094] := 0.1956852;
   Prof_PriceDA.Data[4095] := 0.1956852;
   Prof_PriceDA.Data[4096] := 0.2190564;
   Prof_PriceDA.Data[4097] := 0.2190564;
   Prof_PriceDA.Data[4098] := 0.2190564;
   Prof_PriceDA.Data[4099] := 0.2190564;
   Prof_PriceDA.Data[4100] := 0.3030804;
   Prof_PriceDA.Data[4101] := 0.3030804;
   Prof_PriceDA.Data[4102] := 0.3030804;
   Prof_PriceDA.Data[4103] := 0.3030804;
   Prof_PriceDA.Data[4104] := 0.2873556;
   Prof_PriceDA.Data[4105] := 0.2873556;
   Prof_PriceDA.Data[4106] := 0.2873556;
   Prof_PriceDA.Data[4107] := 0.2873556;
   Prof_PriceDA.Data[4108] := 0.240462;
   Prof_PriceDA.Data[4109] := 0.240462;
   Prof_PriceDA.Data[4110] := 0.240462;
   Prof_PriceDA.Data[4111] := 0.240462;
   Prof_PriceDA.Data[4112] := 0.2384316;
   Prof_PriceDA.Data[4113] := 0.2384316;
   Prof_PriceDA.Data[4114] := 0.2384316;
   Prof_PriceDA.Data[4115] := 0.2384316;
   Prof_PriceDA.Data[4116] := 0.1923156;
   Prof_PriceDA.Data[4117] := 0.1923156;
   Prof_PriceDA.Data[4118] := 0.1923156;
   Prof_PriceDA.Data[4119] := 0.1923156;
   Prof_PriceDA.Data[4120] := 0.1861812;
   Prof_PriceDA.Data[4121] := 0.1861812;
   Prof_PriceDA.Data[4122] := 0.1861812;
   Prof_PriceDA.Data[4123] := 0.1861812;
   Prof_PriceDA.Data[4124] := 0.1728;
   Prof_PriceDA.Data[4125] := 0.1728;
   Prof_PriceDA.Data[4126] := 0.1728;
   Prof_PriceDA.Data[4127] := 0.1728;
   Prof_PriceDA.Data[4128] := 0.1722708;
   Prof_PriceDA.Data[4129] := 0.1722708;
   Prof_PriceDA.Data[4130] := 0.1722708;
   Prof_PriceDA.Data[4131] := 0.1722708;
   Prof_PriceDA.Data[4132] := 0.161298;
   Prof_PriceDA.Data[4133] := 0.161298;
   Prof_PriceDA.Data[4134] := 0.161298;
   Prof_PriceDA.Data[4135] := 0.161298;
   Prof_PriceDA.Data[4136] := 0.158868;
   Prof_PriceDA.Data[4137] := 0.158868;
   Prof_PriceDA.Data[4138] := 0.158868;
   Prof_PriceDA.Data[4139] := 0.158868;
   Prof_PriceDA.Data[4140] := 0.1538136;
   Prof_PriceDA.Data[4141] := 0.1538136;
   Prof_PriceDA.Data[4142] := 0.1538136;
   Prof_PriceDA.Data[4143] := 0.1538136;
   Prof_PriceDA.Data[4144] := 0.1591596;
   Prof_PriceDA.Data[4145] := 0.1591596;
   Prof_PriceDA.Data[4146] := 0.1591596;
   Prof_PriceDA.Data[4147] := 0.1591596;
   Prof_PriceDA.Data[4148] := 0.1767852;
   Prof_PriceDA.Data[4149] := 0.1767852;
   Prof_PriceDA.Data[4150] := 0.1767852;
   Prof_PriceDA.Data[4151] := 0.1767852;
   Prof_PriceDA.Data[4152] := 0.2259684;
   Prof_PriceDA.Data[4153] := 0.2259684;
   Prof_PriceDA.Data[4154] := 0.2259684;
   Prof_PriceDA.Data[4155] := 0.2259684;
   Prof_PriceDA.Data[4156] := 0.421524;
   Prof_PriceDA.Data[4157] := 0.421524;
   Prof_PriceDA.Data[4158] := 0.421524;
   Prof_PriceDA.Data[4159] := 0.421524;
   Prof_PriceDA.Data[4160] := 0.3348108;
   Prof_PriceDA.Data[4161] := 0.3348108;
   Prof_PriceDA.Data[4162] := 0.3348108;
   Prof_PriceDA.Data[4163] := 0.3348108;
   Prof_PriceDA.Data[4164] := 0.2808108;
   Prof_PriceDA.Data[4165] := 0.2808108;
   Prof_PriceDA.Data[4166] := 0.2808108;
   Prof_PriceDA.Data[4167] := 0.2808108;
   Prof_PriceDA.Data[4168] := 0.2247588;
   Prof_PriceDA.Data[4169] := 0.2247588;
   Prof_PriceDA.Data[4170] := 0.2247588;
   Prof_PriceDA.Data[4171] := 0.2247588;
   Prof_PriceDA.Data[4172] := 0.2027268;
   Prof_PriceDA.Data[4173] := 0.2027268;
   Prof_PriceDA.Data[4174] := 0.2027268;
   Prof_PriceDA.Data[4175] := 0.2027268;
   Prof_PriceDA.Data[4176] := 0.2015604;
   Prof_PriceDA.Data[4177] := 0.2015604;
   Prof_PriceDA.Data[4178] := 0.2015604;
   Prof_PriceDA.Data[4179] := 0.2015604;
   Prof_PriceDA.Data[4180] := 0.2252664;
   Prof_PriceDA.Data[4181] := 0.2252664;
   Prof_PriceDA.Data[4182] := 0.2252664;
   Prof_PriceDA.Data[4183] := 0.2252664;
   Prof_PriceDA.Data[4184] := 0.2457648;
   Prof_PriceDA.Data[4185] := 0.2457648;
   Prof_PriceDA.Data[4186] := 0.2457648;
   Prof_PriceDA.Data[4187] := 0.2457648;
   Prof_PriceDA.Data[4188] := 0.2673;
   Prof_PriceDA.Data[4189] := 0.2673;
   Prof_PriceDA.Data[4190] := 0.2673;
   Prof_PriceDA.Data[4191] := 0.2673;
   Prof_PriceDA.Data[4192] := 0.2891484;
   Prof_PriceDA.Data[4193] := 0.2891484;
   Prof_PriceDA.Data[4194] := 0.2891484;
   Prof_PriceDA.Data[4195] := 0.2891484;
   Prof_PriceDA.Data[4196] := 0.2678184;
   Prof_PriceDA.Data[4197] := 0.2678184;
   Prof_PriceDA.Data[4198] := 0.2678184;
   Prof_PriceDA.Data[4199] := 0.2678184;
   Prof_PriceDA.Data[4200] := 0.2236788;
   Prof_PriceDA.Data[4201] := 0.2236788;
   Prof_PriceDA.Data[4202] := 0.2236788;
   Prof_PriceDA.Data[4203] := 0.2236788;
   Prof_PriceDA.Data[4204] := 0.2122416;
   Prof_PriceDA.Data[4205] := 0.2122416;
   Prof_PriceDA.Data[4206] := 0.2122416;
   Prof_PriceDA.Data[4207] := 0.2122416;
   Prof_PriceDA.Data[4208] := 0.1927152;
   Prof_PriceDA.Data[4209] := 0.1927152;
   Prof_PriceDA.Data[4210] := 0.1927152;
   Prof_PriceDA.Data[4211] := 0.1927152;
   Prof_PriceDA.Data[4212] := 0.1759536;
   Prof_PriceDA.Data[4213] := 0.1759536;
   Prof_PriceDA.Data[4214] := 0.1759536;
   Prof_PriceDA.Data[4215] := 0.1759536;
   Prof_PriceDA.Data[4216] := 0.1653696;
   Prof_PriceDA.Data[4217] := 0.1653696;
   Prof_PriceDA.Data[4218] := 0.1653696;
   Prof_PriceDA.Data[4219] := 0.1653696;
   Prof_PriceDA.Data[4220] := 0.1503036;
   Prof_PriceDA.Data[4221] := 0.1503036;
   Prof_PriceDA.Data[4222] := 0.1503036;
   Prof_PriceDA.Data[4223] := 0.1503036;
   Prof_PriceDA.Data[4224] := 0.1514376;
   Prof_PriceDA.Data[4225] := 0.1514376;
   Prof_PriceDA.Data[4226] := 0.1514376;
   Prof_PriceDA.Data[4227] := 0.1514376;
   Prof_PriceDA.Data[4228] := 0.1460916;
   Prof_PriceDA.Data[4229] := 0.1460916;
   Prof_PriceDA.Data[4230] := 0.1460916;
   Prof_PriceDA.Data[4231] := 0.1460916;
   Prof_PriceDA.Data[4232] := 0.141048;
   Prof_PriceDA.Data[4233] := 0.141048;
   Prof_PriceDA.Data[4234] := 0.141048;
   Prof_PriceDA.Data[4235] := 0.141048;
   Prof_PriceDA.Data[4236] := 0.1412748;
   Prof_PriceDA.Data[4237] := 0.1412748;
   Prof_PriceDA.Data[4238] := 0.1412748;
   Prof_PriceDA.Data[4239] := 0.1412748;
   Prof_PriceDA.Data[4240] := 0.141858;
   Prof_PriceDA.Data[4241] := 0.141858;
   Prof_PriceDA.Data[4242] := 0.141858;
   Prof_PriceDA.Data[4243] := 0.141858;
   Prof_PriceDA.Data[4244] := 0.1520748;
   Prof_PriceDA.Data[4245] := 0.1520748;
   Prof_PriceDA.Data[4246] := 0.1520748;
   Prof_PriceDA.Data[4247] := 0.1520748;
   Prof_PriceDA.Data[4248] := 0.1772712;
   Prof_PriceDA.Data[4249] := 0.1772712;
   Prof_PriceDA.Data[4250] := 0.1772712;
   Prof_PriceDA.Data[4251] := 0.1772712;
   Prof_PriceDA.Data[4252] := 0.2337336;
   Prof_PriceDA.Data[4253] := 0.2337336;
   Prof_PriceDA.Data[4254] := 0.2337336;
   Prof_PriceDA.Data[4255] := 0.2337336;
   Prof_PriceDA.Data[4256] := 0.2835216;
   Prof_PriceDA.Data[4257] := 0.2835216;
   Prof_PriceDA.Data[4258] := 0.2835216;
   Prof_PriceDA.Data[4259] := 0.2835216;
   Prof_PriceDA.Data[4260] := 0.229284;
   Prof_PriceDA.Data[4261] := 0.229284;
   Prof_PriceDA.Data[4262] := 0.229284;
   Prof_PriceDA.Data[4263] := 0.229284;
   Prof_PriceDA.Data[4264] := 0.1935144;
   Prof_PriceDA.Data[4265] := 0.1935144;
   Prof_PriceDA.Data[4266] := 0.1935144;
   Prof_PriceDA.Data[4267] := 0.1935144;
   Prof_PriceDA.Data[4268] := 0.1778976;
   Prof_PriceDA.Data[4269] := 0.1778976;
   Prof_PriceDA.Data[4270] := 0.1778976;
   Prof_PriceDA.Data[4271] := 0.1778976;
   Prof_PriceDA.Data[4272] := 0.1623564;
   Prof_PriceDA.Data[4273] := 0.1623564;
   Prof_PriceDA.Data[4274] := 0.1623564;
   Prof_PriceDA.Data[4275] := 0.1623564;
   Prof_PriceDA.Data[4276] := 0.1625508;
   Prof_PriceDA.Data[4277] := 0.1625508;
   Prof_PriceDA.Data[4278] := 0.1625508;
   Prof_PriceDA.Data[4279] := 0.1625508;
   Prof_PriceDA.Data[4280] := 0.1714824;
   Prof_PriceDA.Data[4281] := 0.1714824;
   Prof_PriceDA.Data[4282] := 0.1714824;
   Prof_PriceDA.Data[4283] := 0.1714824;
   Prof_PriceDA.Data[4284] := 0.1871316;
   Prof_PriceDA.Data[4285] := 0.1871316;
   Prof_PriceDA.Data[4286] := 0.1871316;
   Prof_PriceDA.Data[4287] := 0.1871316;
   Prof_PriceDA.Data[4288] := 0.2142396;
   Prof_PriceDA.Data[4289] := 0.2142396;
   Prof_PriceDA.Data[4290] := 0.2142396;
   Prof_PriceDA.Data[4291] := 0.2142396;
   Prof_PriceDA.Data[4292] := 0.3135456;
   Prof_PriceDA.Data[4293] := 0.3135456;
   Prof_PriceDA.Data[4294] := 0.3135456;
   Prof_PriceDA.Data[4295] := 0.3135456;
   Prof_PriceDA.Data[4296] := 0.3104244;
   Prof_PriceDA.Data[4297] := 0.3104244;
   Prof_PriceDA.Data[4298] := 0.3104244;
   Prof_PriceDA.Data[4299] := 0.3104244;
   Prof_PriceDA.Data[4300] := 0.2420388;
   Prof_PriceDA.Data[4301] := 0.2420388;
   Prof_PriceDA.Data[4302] := 0.2420388;
   Prof_PriceDA.Data[4303] := 0.2420388;
   Prof_PriceDA.Data[4304] := 0.198234;
   Prof_PriceDA.Data[4305] := 0.198234;
   Prof_PriceDA.Data[4306] := 0.198234;
   Prof_PriceDA.Data[4307] := 0.198234;
   Prof_PriceDA.Data[4308] := 0.1766232;
   Prof_PriceDA.Data[4309] := 0.1766232;
   Prof_PriceDA.Data[4310] := 0.1766232;
   Prof_PriceDA.Data[4311] := 0.1766232;
   Prof_PriceDA.Data[4312] := 0.16524;
   Prof_PriceDA.Data[4313] := 0.16524;
   Prof_PriceDA.Data[4314] := 0.16524;
   Prof_PriceDA.Data[4315] := 0.16524;
   Prof_PriceDA.Data[4316] := 0.1512324;
   Prof_PriceDA.Data[4317] := 0.1512324;
   Prof_PriceDA.Data[4318] := 0.1512324;
   Prof_PriceDA.Data[4319] := 0.1512324;
   Prof_PriceDA.Data[4320] := 0.1472688;
   Prof_PriceDA.Data[4321] := 0.1472688;
   Prof_PriceDA.Data[4322] := 0.1472688;
   Prof_PriceDA.Data[4323] := 0.1472688;
   Prof_PriceDA.Data[4324] := 0.1418796;
   Prof_PriceDA.Data[4325] := 0.1418796;
   Prof_PriceDA.Data[4326] := 0.1418796;
   Prof_PriceDA.Data[4327] := 0.1418796;
   Prof_PriceDA.Data[4328] := 0.1303884;
   Prof_PriceDA.Data[4329] := 0.1303884;
   Prof_PriceDA.Data[4330] := 0.1303884;
   Prof_PriceDA.Data[4331] := 0.1303884;
   Prof_PriceDA.Data[4332] := 0.1291356;
   Prof_PriceDA.Data[4333] := 0.1291356;
   Prof_PriceDA.Data[4334] := 0.1291356;
   Prof_PriceDA.Data[4335] := 0.1291356;
   Prof_PriceDA.Data[4336] := 0.1295784;
   Prof_PriceDA.Data[4337] := 0.1295784;
   Prof_PriceDA.Data[4338] := 0.1295784;
   Prof_PriceDA.Data[4339] := 0.1295784;
   Prof_PriceDA.Data[4340] := 0.1315872;
   Prof_PriceDA.Data[4341] := 0.1315872;
   Prof_PriceDA.Data[4342] := 0.1315872;
   Prof_PriceDA.Data[4343] := 0.1315872;
   Prof_PriceDA.Data[4344] := 0.146718;
   Prof_PriceDA.Data[4345] := 0.146718;
   Prof_PriceDA.Data[4346] := 0.146718;
   Prof_PriceDA.Data[4347] := 0.146718;
   Prof_PriceDA.Data[4348] := 0.1623888;
   Prof_PriceDA.Data[4349] := 0.1623888;
   Prof_PriceDA.Data[4350] := 0.1623888;
   Prof_PriceDA.Data[4351] := 0.1623888;
   Prof_PriceDA.Data[4352] := 0.1616328;
   Prof_PriceDA.Data[4353] := 0.1616328;
   Prof_PriceDA.Data[4354] := 0.1616328;
   Prof_PriceDA.Data[4355] := 0.1616328;
   Prof_PriceDA.Data[4356] := 0.148068;
   Prof_PriceDA.Data[4357] := 0.148068;
   Prof_PriceDA.Data[4358] := 0.148068;
   Prof_PriceDA.Data[4359] := 0.148068;
   Prof_PriceDA.Data[4360] := 0.1345572;
   Prof_PriceDA.Data[4361] := 0.1345572;
   Prof_PriceDA.Data[4362] := 0.1345572;
   Prof_PriceDA.Data[4363] := 0.1345572;
   Prof_PriceDA.Data[4364] := 0.1278288;
   Prof_PriceDA.Data[4365] := 0.1278288;
   Prof_PriceDA.Data[4366] := 0.1278288;
   Prof_PriceDA.Data[4367] := 0.1278288;
   Prof_PriceDA.Data[4368] := 0.1213812;
   Prof_PriceDA.Data[4369] := 0.1213812;
   Prof_PriceDA.Data[4370] := 0.1213812;
   Prof_PriceDA.Data[4371] := 0.1213812;
   Prof_PriceDA.Data[4372] := 0.1188108;
   Prof_PriceDA.Data[4373] := 0.1188108;
   Prof_PriceDA.Data[4374] := 0.1188108;
   Prof_PriceDA.Data[4375] := 0.1188108;
   Prof_PriceDA.Data[4376] := 0.126252;
   Prof_PriceDA.Data[4377] := 0.126252;
   Prof_PriceDA.Data[4378] := 0.126252;
   Prof_PriceDA.Data[4379] := 0.126252;
   Prof_PriceDA.Data[4380] := 0.1413936;
   Prof_PriceDA.Data[4381] := 0.1413936;
   Prof_PriceDA.Data[4382] := 0.1413936;
   Prof_PriceDA.Data[4383] := 0.1413936;
   Prof_PriceDA.Data[4384] := 0.1687716;
   Prof_PriceDA.Data[4385] := 0.1687716;
   Prof_PriceDA.Data[4386] := 0.1687716;
   Prof_PriceDA.Data[4387] := 0.1687716;
   Prof_PriceDA.Data[4388] := 0.1905552;
   Prof_PriceDA.Data[4389] := 0.1905552;
   Prof_PriceDA.Data[4390] := 0.1905552;
   Prof_PriceDA.Data[4391] := 0.1905552;
   Prof_PriceDA.Data[4392] := 0.1925856;
   Prof_PriceDA.Data[4393] := 0.1925856;
   Prof_PriceDA.Data[4394] := 0.1925856;
   Prof_PriceDA.Data[4395] := 0.1925856;
   Prof_PriceDA.Data[4396] := 0.1880064;
   Prof_PriceDA.Data[4397] := 0.1880064;
   Prof_PriceDA.Data[4398] := 0.1880064;
   Prof_PriceDA.Data[4399] := 0.1880064;
   Prof_PriceDA.Data[4400] := 0.1818504;
   Prof_PriceDA.Data[4401] := 0.1818504;
   Prof_PriceDA.Data[4402] := 0.1818504;
   Prof_PriceDA.Data[4403] := 0.1818504;
   Prof_PriceDA.Data[4404] := 0.165348;
   Prof_PriceDA.Data[4405] := 0.165348;
   Prof_PriceDA.Data[4406] := 0.165348;
   Prof_PriceDA.Data[4407] := 0.165348;
   Prof_PriceDA.Data[4408] := 0.1515672;
   Prof_PriceDA.Data[4409] := 0.1515672;
   Prof_PriceDA.Data[4410] := 0.1515672;
   Prof_PriceDA.Data[4411] := 0.1515672;
   Prof_PriceDA.Data[4412] := 0.1441692;
   Prof_PriceDA.Data[4413] := 0.1441692;
   Prof_PriceDA.Data[4414] := 0.1441692;
   Prof_PriceDA.Data[4415] := 0.1441692;
   Prof_PriceDA.Data[4416] := 0.1448388;
   Prof_PriceDA.Data[4417] := 0.1448388;
   Prof_PriceDA.Data[4418] := 0.1448388;
   Prof_PriceDA.Data[4419] := 0.1448388;
   Prof_PriceDA.Data[4420] := 0.139212;
   Prof_PriceDA.Data[4421] := 0.139212;
   Prof_PriceDA.Data[4422] := 0.139212;
   Prof_PriceDA.Data[4423] := 0.139212;
   Prof_PriceDA.Data[4424] := 0.1334556;
   Prof_PriceDA.Data[4425] := 0.1334556;
   Prof_PriceDA.Data[4426] := 0.1334556;
   Prof_PriceDA.Data[4427] := 0.1334556;
   Prof_PriceDA.Data[4428] := 0.129492;
   Prof_PriceDA.Data[4429] := 0.129492;
   Prof_PriceDA.Data[4430] := 0.129492;
   Prof_PriceDA.Data[4431] := 0.129492;
   Prof_PriceDA.Data[4432] := 0.1291356;
   Prof_PriceDA.Data[4433] := 0.1291356;
   Prof_PriceDA.Data[4434] := 0.1291356;
   Prof_PriceDA.Data[4435] := 0.1291356;
   Prof_PriceDA.Data[4436] := 0.1305612;
   Prof_PriceDA.Data[4437] := 0.1305612;
   Prof_PriceDA.Data[4438] := 0.1305612;
   Prof_PriceDA.Data[4439] := 0.1305612;
   Prof_PriceDA.Data[4440] := 0.133758;
   Prof_PriceDA.Data[4441] := 0.133758;
   Prof_PriceDA.Data[4442] := 0.133758;
   Prof_PriceDA.Data[4443] := 0.133758;
   Prof_PriceDA.Data[4444] := 0.1448712;
   Prof_PriceDA.Data[4445] := 0.1448712;
   Prof_PriceDA.Data[4446] := 0.1448712;
   Prof_PriceDA.Data[4447] := 0.1448712;
   Prof_PriceDA.Data[4448] := 0.153846;
   Prof_PriceDA.Data[4449] := 0.153846;
   Prof_PriceDA.Data[4450] := 0.153846;
   Prof_PriceDA.Data[4451] := 0.153846;
   Prof_PriceDA.Data[4452] := 0.152334;
   Prof_PriceDA.Data[4453] := 0.152334;
   Prof_PriceDA.Data[4454] := 0.152334;
   Prof_PriceDA.Data[4455] := 0.152334;
   Prof_PriceDA.Data[4456] := 0.1427652;
   Prof_PriceDA.Data[4457] := 0.1427652;
   Prof_PriceDA.Data[4458] := 0.1427652;
   Prof_PriceDA.Data[4459] := 0.1427652;
   Prof_PriceDA.Data[4460] := 0.141696;
   Prof_PriceDA.Data[4461] := 0.141696;
   Prof_PriceDA.Data[4462] := 0.141696;
   Prof_PriceDA.Data[4463] := 0.141696;
   Prof_PriceDA.Data[4464] := 0.1389636;
   Prof_PriceDA.Data[4465] := 0.1389636;
   Prof_PriceDA.Data[4466] := 0.1389636;
   Prof_PriceDA.Data[4467] := 0.1389636;
   Prof_PriceDA.Data[4468] := 0.1375812;
   Prof_PriceDA.Data[4469] := 0.1375812;
   Prof_PriceDA.Data[4470] := 0.1375812;
   Prof_PriceDA.Data[4471] := 0.1375812;
   Prof_PriceDA.Data[4472] := 0.14094;
   Prof_PriceDA.Data[4473] := 0.14094;
   Prof_PriceDA.Data[4474] := 0.14094;
   Prof_PriceDA.Data[4475] := 0.14094;
   Prof_PriceDA.Data[4476] := 0.1524744;
   Prof_PriceDA.Data[4477] := 0.1524744;
   Prof_PriceDA.Data[4478] := 0.1524744;
   Prof_PriceDA.Data[4479] := 0.1524744;
   Prof_PriceDA.Data[4480] := 0.174852;
   Prof_PriceDA.Data[4481] := 0.174852;
   Prof_PriceDA.Data[4482] := 0.174852;
   Prof_PriceDA.Data[4483] := 0.174852;
   Prof_PriceDA.Data[4484] := 0.1890324;
   Prof_PriceDA.Data[4485] := 0.1890324;
   Prof_PriceDA.Data[4486] := 0.1890324;
   Prof_PriceDA.Data[4487] := 0.1890324;
   Prof_PriceDA.Data[4488] := 0.191322;
   Prof_PriceDA.Data[4489] := 0.191322;
   Prof_PriceDA.Data[4490] := 0.191322;
   Prof_PriceDA.Data[4491] := 0.191322;
   Prof_PriceDA.Data[4492] := 0.1876932;
   Prof_PriceDA.Data[4493] := 0.1876932;
   Prof_PriceDA.Data[4494] := 0.1876932;
   Prof_PriceDA.Data[4495] := 0.1876932;
   Prof_PriceDA.Data[4496] := 0.1830708;
   Prof_PriceDA.Data[4497] := 0.1830708;
   Prof_PriceDA.Data[4498] := 0.1830708;
   Prof_PriceDA.Data[4499] := 0.1830708;
   Prof_PriceDA.Data[4500] := 0.1726272;
   Prof_PriceDA.Data[4501] := 0.1726272;
   Prof_PriceDA.Data[4502] := 0.1726272;
   Prof_PriceDA.Data[4503] := 0.1726272;
   Prof_PriceDA.Data[4504] := 0.1613412;
   Prof_PriceDA.Data[4505] := 0.1613412;
   Prof_PriceDA.Data[4506] := 0.1613412;
   Prof_PriceDA.Data[4507] := 0.1613412;
   Prof_PriceDA.Data[4508] := 0.1420308;
   Prof_PriceDA.Data[4509] := 0.1420308;
   Prof_PriceDA.Data[4510] := 0.1420308;
   Prof_PriceDA.Data[4511] := 0.1420308;
   Prof_PriceDA.Data[4512] := 0.1431216;
   Prof_PriceDA.Data[4513] := 0.1431216;
   Prof_PriceDA.Data[4514] := 0.1431216;
   Prof_PriceDA.Data[4515] := 0.1431216;
   Prof_PriceDA.Data[4516] := 0.1307448;
   Prof_PriceDA.Data[4517] := 0.1307448;
   Prof_PriceDA.Data[4518] := 0.1307448;
   Prof_PriceDA.Data[4519] := 0.1307448;
   Prof_PriceDA.Data[4520] := 0.1299672;
   Prof_PriceDA.Data[4521] := 0.1299672;
   Prof_PriceDA.Data[4522] := 0.1299672;
   Prof_PriceDA.Data[4523] := 0.1299672;
   Prof_PriceDA.Data[4524] := 0.1365876;
   Prof_PriceDA.Data[4525] := 0.1365876;
   Prof_PriceDA.Data[4526] := 0.1365876;
   Prof_PriceDA.Data[4527] := 0.1365876;
   Prof_PriceDA.Data[4528] := 0.1406052;
   Prof_PriceDA.Data[4529] := 0.1406052;
   Prof_PriceDA.Data[4530] := 0.1406052;
   Prof_PriceDA.Data[4531] := 0.1406052;
   Prof_PriceDA.Data[4532] := 0.1550124;
   Prof_PriceDA.Data[4533] := 0.1550124;
   Prof_PriceDA.Data[4534] := 0.1550124;
   Prof_PriceDA.Data[4535] := 0.1550124;
   Prof_PriceDA.Data[4536] := 0.1884924;
   Prof_PriceDA.Data[4537] := 0.1884924;
   Prof_PriceDA.Data[4538] := 0.1884924;
   Prof_PriceDA.Data[4539] := 0.1884924;
   Prof_PriceDA.Data[4540] := 0.2253096;
   Prof_PriceDA.Data[4541] := 0.2253096;
   Prof_PriceDA.Data[4542] := 0.2253096;
   Prof_PriceDA.Data[4543] := 0.2253096;
   Prof_PriceDA.Data[4544] := 0.2265732;
   Prof_PriceDA.Data[4545] := 0.2265732;
   Prof_PriceDA.Data[4546] := 0.2265732;
   Prof_PriceDA.Data[4547] := 0.2265732;
   Prof_PriceDA.Data[4548] := 0.185004;
   Prof_PriceDA.Data[4549] := 0.185004;
   Prof_PriceDA.Data[4550] := 0.185004;
   Prof_PriceDA.Data[4551] := 0.185004;
   Prof_PriceDA.Data[4552] := 0.1508436;
   Prof_PriceDA.Data[4553] := 0.1508436;
   Prof_PriceDA.Data[4554] := 0.1508436;
   Prof_PriceDA.Data[4555] := 0.1508436;
   Prof_PriceDA.Data[4556] := 0.1288764;
   Prof_PriceDA.Data[4557] := 0.1288764;
   Prof_PriceDA.Data[4558] := 0.1288764;
   Prof_PriceDA.Data[4559] := 0.1288764;
   Prof_PriceDA.Data[4560] := 0.1232928;
   Prof_PriceDA.Data[4561] := 0.1232928;
   Prof_PriceDA.Data[4562] := 0.1232928;
   Prof_PriceDA.Data[4563] := 0.1232928;
   Prof_PriceDA.Data[4564] := 0.1176012;
   Prof_PriceDA.Data[4565] := 0.1176012;
   Prof_PriceDA.Data[4566] := 0.1176012;
   Prof_PriceDA.Data[4567] := 0.1176012;
   Prof_PriceDA.Data[4568] := 0.13176;
   Prof_PriceDA.Data[4569] := 0.13176;
   Prof_PriceDA.Data[4570] := 0.13176;
   Prof_PriceDA.Data[4571] := 0.13176;
   Prof_PriceDA.Data[4572] := 0.1601748;
   Prof_PriceDA.Data[4573] := 0.1601748;
   Prof_PriceDA.Data[4574] := 0.1601748;
   Prof_PriceDA.Data[4575] := 0.1601748;
   Prof_PriceDA.Data[4576] := 0.1869372;
   Prof_PriceDA.Data[4577] := 0.1869372;
   Prof_PriceDA.Data[4578] := 0.1869372;
   Prof_PriceDA.Data[4579] := 0.1869372;
   Prof_PriceDA.Data[4580] := 0.238572;
   Prof_PriceDA.Data[4581] := 0.238572;
   Prof_PriceDA.Data[4582] := 0.238572;
   Prof_PriceDA.Data[4583] := 0.238572;
   Prof_PriceDA.Data[4584] := 0.2883816;
   Prof_PriceDA.Data[4585] := 0.2883816;
   Prof_PriceDA.Data[4586] := 0.2883816;
   Prof_PriceDA.Data[4587] := 0.2883816;
   Prof_PriceDA.Data[4588] := 0.2338956;
   Prof_PriceDA.Data[4589] := 0.2338956;
   Prof_PriceDA.Data[4590] := 0.2338956;
   Prof_PriceDA.Data[4591] := 0.2338956;
   Prof_PriceDA.Data[4592] := 0.1934928;
   Prof_PriceDA.Data[4593] := 0.1934928;
   Prof_PriceDA.Data[4594] := 0.1934928;
   Prof_PriceDA.Data[4595] := 0.1934928;
   Prof_PriceDA.Data[4596] := 0.1759212;
   Prof_PriceDA.Data[4597] := 0.1759212;
   Prof_PriceDA.Data[4598] := 0.1759212;
   Prof_PriceDA.Data[4599] := 0.1759212;
   Prof_PriceDA.Data[4600] := 0.169074;
   Prof_PriceDA.Data[4601] := 0.169074;
   Prof_PriceDA.Data[4602] := 0.169074;
   Prof_PriceDA.Data[4603] := 0.169074;
   Prof_PriceDA.Data[4604] := 0.15444;
   Prof_PriceDA.Data[4605] := 0.15444;
   Prof_PriceDA.Data[4606] := 0.15444;
   Prof_PriceDA.Data[4607] := 0.15444;
   Prof_PriceDA.Data[4608] := 0.146664;
   Prof_PriceDA.Data[4609] := 0.146664;
   Prof_PriceDA.Data[4610] := 0.146664;
   Prof_PriceDA.Data[4611] := 0.146664;
   Prof_PriceDA.Data[4612] := 0.1429488;
   Prof_PriceDA.Data[4613] := 0.1429488;
   Prof_PriceDA.Data[4614] := 0.1429488;
   Prof_PriceDA.Data[4615] := 0.1429488;
   Prof_PriceDA.Data[4616] := 0.1358748;
   Prof_PriceDA.Data[4617] := 0.1358748;
   Prof_PriceDA.Data[4618] := 0.1358748;
   Prof_PriceDA.Data[4619] := 0.1358748;
   Prof_PriceDA.Data[4620] := 0.1331316;
   Prof_PriceDA.Data[4621] := 0.1331316;
   Prof_PriceDA.Data[4622] := 0.1331316;
   Prof_PriceDA.Data[4623] := 0.1331316;
   Prof_PriceDA.Data[4624] := 0.1377216;
   Prof_PriceDA.Data[4625] := 0.1377216;
   Prof_PriceDA.Data[4626] := 0.1377216;
   Prof_PriceDA.Data[4627] := 0.1377216;
   Prof_PriceDA.Data[4628] := 0.163998;
   Prof_PriceDA.Data[4629] := 0.163998;
   Prof_PriceDA.Data[4630] := 0.163998;
   Prof_PriceDA.Data[4631] := 0.163998;
   Prof_PriceDA.Data[4632] := 0.2263032;
   Prof_PriceDA.Data[4633] := 0.2263032;
   Prof_PriceDA.Data[4634] := 0.2263032;
   Prof_PriceDA.Data[4635] := 0.2263032;
   Prof_PriceDA.Data[4636] := 0.3576096;
   Prof_PriceDA.Data[4637] := 0.3576096;
   Prof_PriceDA.Data[4638] := 0.3576096;
   Prof_PriceDA.Data[4639] := 0.3576096;
   Prof_PriceDA.Data[4640] := 0.209304;
   Prof_PriceDA.Data[4641] := 0.209304;
   Prof_PriceDA.Data[4642] := 0.209304;
   Prof_PriceDA.Data[4643] := 0.209304;
   Prof_PriceDA.Data[4644] := 0.1750356;
   Prof_PriceDA.Data[4645] := 0.1750356;
   Prof_PriceDA.Data[4646] := 0.1750356;
   Prof_PriceDA.Data[4647] := 0.1750356;
   Prof_PriceDA.Data[4648] := 0.154386;
   Prof_PriceDA.Data[4649] := 0.154386;
   Prof_PriceDA.Data[4650] := 0.154386;
   Prof_PriceDA.Data[4651] := 0.154386;
   Prof_PriceDA.Data[4652] := 0.1445148;
   Prof_PriceDA.Data[4653] := 0.1445148;
   Prof_PriceDA.Data[4654] := 0.1445148;
   Prof_PriceDA.Data[4655] := 0.1445148;
   Prof_PriceDA.Data[4656] := 0.142398;
   Prof_PriceDA.Data[4657] := 0.142398;
   Prof_PriceDA.Data[4658] := 0.142398;
   Prof_PriceDA.Data[4659] := 0.142398;
   Prof_PriceDA.Data[4660] := 0.1559736;
   Prof_PriceDA.Data[4661] := 0.1559736;
   Prof_PriceDA.Data[4662] := 0.1559736;
   Prof_PriceDA.Data[4663] := 0.1559736;
   Prof_PriceDA.Data[4664] := 0.1631448;
   Prof_PriceDA.Data[4665] := 0.1631448;
   Prof_PriceDA.Data[4666] := 0.1631448;
   Prof_PriceDA.Data[4667] := 0.1631448;
   Prof_PriceDA.Data[4668] := 0.1770876;
   Prof_PriceDA.Data[4669] := 0.1770876;
   Prof_PriceDA.Data[4670] := 0.1770876;
   Prof_PriceDA.Data[4671] := 0.1770876;
   Prof_PriceDA.Data[4672] := 0.3453516;
   Prof_PriceDA.Data[4673] := 0.3453516;
   Prof_PriceDA.Data[4674] := 0.3453516;
   Prof_PriceDA.Data[4675] := 0.3453516;
   Prof_PriceDA.Data[4676] := 0.2810268;
   Prof_PriceDA.Data[4677] := 0.2810268;
   Prof_PriceDA.Data[4678] := 0.2810268;
   Prof_PriceDA.Data[4679] := 0.2810268;
   Prof_PriceDA.Data[4680] := 0.2770092;
   Prof_PriceDA.Data[4681] := 0.2770092;
   Prof_PriceDA.Data[4682] := 0.2770092;
   Prof_PriceDA.Data[4683] := 0.2770092;
   Prof_PriceDA.Data[4684] := 0.2601612;
   Prof_PriceDA.Data[4685] := 0.2601612;
   Prof_PriceDA.Data[4686] := 0.2601612;
   Prof_PriceDA.Data[4687] := 0.2601612;
   Prof_PriceDA.Data[4688] := 0.1939248;
   Prof_PriceDA.Data[4689] := 0.1939248;
   Prof_PriceDA.Data[4690] := 0.1939248;
   Prof_PriceDA.Data[4691] := 0.1939248;
   Prof_PriceDA.Data[4692] := 0.1817316;
   Prof_PriceDA.Data[4693] := 0.1817316;
   Prof_PriceDA.Data[4694] := 0.1817316;
   Prof_PriceDA.Data[4695] := 0.1817316;
   Prof_PriceDA.Data[4696] := 0.1740852;
   Prof_PriceDA.Data[4697] := 0.1740852;
   Prof_PriceDA.Data[4698] := 0.1740852;
   Prof_PriceDA.Data[4699] := 0.1740852;
   Prof_PriceDA.Data[4700] := 0.1480032;
   Prof_PriceDA.Data[4701] := 0.1480032;
   Prof_PriceDA.Data[4702] := 0.1480032;
   Prof_PriceDA.Data[4703] := 0.1480032;
   Prof_PriceDA.Data[4704] := 0.14121;
   Prof_PriceDA.Data[4705] := 0.14121;
   Prof_PriceDA.Data[4706] := 0.14121;
   Prof_PriceDA.Data[4707] := 0.14121;
   Prof_PriceDA.Data[4708] := 0.1392768;
   Prof_PriceDA.Data[4709] := 0.1392768;
   Prof_PriceDA.Data[4710] := 0.1392768;
   Prof_PriceDA.Data[4711] := 0.1392768;
   Prof_PriceDA.Data[4712] := 0.1372896;
   Prof_PriceDA.Data[4713] := 0.1372896;
   Prof_PriceDA.Data[4714] := 0.1372896;
   Prof_PriceDA.Data[4715] := 0.1372896;
   Prof_PriceDA.Data[4716] := 0.136458;
   Prof_PriceDA.Data[4717] := 0.136458;
   Prof_PriceDA.Data[4718] := 0.136458;
   Prof_PriceDA.Data[4719] := 0.136458;
   Prof_PriceDA.Data[4720] := 0.1398168;
   Prof_PriceDA.Data[4721] := 0.1398168;
   Prof_PriceDA.Data[4722] := 0.1398168;
   Prof_PriceDA.Data[4723] := 0.1398168;
   Prof_PriceDA.Data[4724] := 0.155088;
   Prof_PriceDA.Data[4725] := 0.155088;
   Prof_PriceDA.Data[4726] := 0.155088;
   Prof_PriceDA.Data[4727] := 0.155088;
   Prof_PriceDA.Data[4728] := 0.1828872;
   Prof_PriceDA.Data[4729] := 0.1828872;
   Prof_PriceDA.Data[4730] := 0.1828872;
   Prof_PriceDA.Data[4731] := 0.1828872;
   Prof_PriceDA.Data[4732] := 0.218592;
   Prof_PriceDA.Data[4733] := 0.218592;
   Prof_PriceDA.Data[4734] := 0.218592;
   Prof_PriceDA.Data[4735] := 0.218592;
   Prof_PriceDA.Data[4736] := 0.190404;
   Prof_PriceDA.Data[4737] := 0.190404;
   Prof_PriceDA.Data[4738] := 0.190404;
   Prof_PriceDA.Data[4739] := 0.190404;
   Prof_PriceDA.Data[4740] := 0.165456;
   Prof_PriceDA.Data[4741] := 0.165456;
   Prof_PriceDA.Data[4742] := 0.165456;
   Prof_PriceDA.Data[4743] := 0.165456;
   Prof_PriceDA.Data[4744] := 0.123606;
   Prof_PriceDA.Data[4745] := 0.123606;
   Prof_PriceDA.Data[4746] := 0.123606;
   Prof_PriceDA.Data[4747] := 0.123606;
   Prof_PriceDA.Data[4748] := 0.1240056;
   Prof_PriceDA.Data[4749] := 0.1240056;
   Prof_PriceDA.Data[4750] := 0.1240056;
   Prof_PriceDA.Data[4751] := 0.1240056;
   Prof_PriceDA.Data[4752] := 0.1162728;
   Prof_PriceDA.Data[4753] := 0.1162728;
   Prof_PriceDA.Data[4754] := 0.1162728;
   Prof_PriceDA.Data[4755] := 0.1162728;
   Prof_PriceDA.Data[4756] := 0.1160568;
   Prof_PriceDA.Data[4757] := 0.1160568;
   Prof_PriceDA.Data[4758] := 0.1160568;
   Prof_PriceDA.Data[4759] := 0.1160568;
   Prof_PriceDA.Data[4760] := 0.126954;
   Prof_PriceDA.Data[4761] := 0.126954;
   Prof_PriceDA.Data[4762] := 0.126954;
   Prof_PriceDA.Data[4763] := 0.126954;
   Prof_PriceDA.Data[4764] := 0.1515888;
   Prof_PriceDA.Data[4765] := 0.1515888;
   Prof_PriceDA.Data[4766] := 0.1515888;
   Prof_PriceDA.Data[4767] := 0.1515888;
   Prof_PriceDA.Data[4768] := 0.190944;
   Prof_PriceDA.Data[4769] := 0.190944;
   Prof_PriceDA.Data[4770] := 0.190944;
   Prof_PriceDA.Data[4771] := 0.190944;
   Prof_PriceDA.Data[4772] := 0.249534;
   Prof_PriceDA.Data[4773] := 0.249534;
   Prof_PriceDA.Data[4774] := 0.249534;
   Prof_PriceDA.Data[4775] := 0.249534;
   Prof_PriceDA.Data[4776] := 0.2520504;
   Prof_PriceDA.Data[4777] := 0.2520504;
   Prof_PriceDA.Data[4778] := 0.2520504;
   Prof_PriceDA.Data[4779] := 0.2520504;
   Prof_PriceDA.Data[4780] := 0.2164968;
   Prof_PriceDA.Data[4781] := 0.2164968;
   Prof_PriceDA.Data[4782] := 0.2164968;
   Prof_PriceDA.Data[4783] := 0.2164968;
   Prof_PriceDA.Data[4784] := 0.1938492;
   Prof_PriceDA.Data[4785] := 0.1938492;
   Prof_PriceDA.Data[4786] := 0.1938492;
   Prof_PriceDA.Data[4787] := 0.1938492;
   Prof_PriceDA.Data[4788] := 0.1805868;
   Prof_PriceDA.Data[4789] := 0.1805868;
   Prof_PriceDA.Data[4790] := 0.1805868;
   Prof_PriceDA.Data[4791] := 0.1805868;
   Prof_PriceDA.Data[4792] := 0.1764936;
   Prof_PriceDA.Data[4793] := 0.1764936;
   Prof_PriceDA.Data[4794] := 0.1764936;
   Prof_PriceDA.Data[4795] := 0.1764936;
   Prof_PriceDA.Data[4796] := 0.1671192;
   Prof_PriceDA.Data[4797] := 0.1671192;
   Prof_PriceDA.Data[4798] := 0.1671192;
   Prof_PriceDA.Data[4799] := 0.1671192;
   Prof_PriceDA.Data[4800] := 0.1350972;
   Prof_PriceDA.Data[4801] := 0.1350972;
   Prof_PriceDA.Data[4802] := 0.1350972;
   Prof_PriceDA.Data[4803] := 0.1350972;
   Prof_PriceDA.Data[4804] := 0.1303452;
   Prof_PriceDA.Data[4805] := 0.1303452;
   Prof_PriceDA.Data[4806] := 0.1303452;
   Prof_PriceDA.Data[4807] := 0.1303452;
   Prof_PriceDA.Data[4808] := 0.1251936;
   Prof_PriceDA.Data[4809] := 0.1251936;
   Prof_PriceDA.Data[4810] := 0.1251936;
   Prof_PriceDA.Data[4811] := 0.1251936;
   Prof_PriceDA.Data[4812] := 0.1203984;
   Prof_PriceDA.Data[4813] := 0.1203984;
   Prof_PriceDA.Data[4814] := 0.1203984;
   Prof_PriceDA.Data[4815] := 0.1203984;
   Prof_PriceDA.Data[4816] := 0.1305396;
   Prof_PriceDA.Data[4817] := 0.1305396;
   Prof_PriceDA.Data[4818] := 0.1305396;
   Prof_PriceDA.Data[4819] := 0.1305396;
   Prof_PriceDA.Data[4820] := 0.1563948;
   Prof_PriceDA.Data[4821] := 0.1563948;
   Prof_PriceDA.Data[4822] := 0.1563948;
   Prof_PriceDA.Data[4823] := 0.1563948;
   Prof_PriceDA.Data[4824] := 0.2001456;
   Prof_PriceDA.Data[4825] := 0.2001456;
   Prof_PriceDA.Data[4826] := 0.2001456;
   Prof_PriceDA.Data[4827] := 0.2001456;
   Prof_PriceDA.Data[4828] := 0.263412;
   Prof_PriceDA.Data[4829] := 0.263412;
   Prof_PriceDA.Data[4830] := 0.263412;
   Prof_PriceDA.Data[4831] := 0.263412;
   Prof_PriceDA.Data[4832] := 0.19062;
   Prof_PriceDA.Data[4833] := 0.19062;
   Prof_PriceDA.Data[4834] := 0.19062;
   Prof_PriceDA.Data[4835] := 0.19062;
   Prof_PriceDA.Data[4836] := 0.1302804;
   Prof_PriceDA.Data[4837] := 0.1302804;
   Prof_PriceDA.Data[4838] := 0.1302804;
   Prof_PriceDA.Data[4839] := 0.1302804;
   Prof_PriceDA.Data[4840] := 0.1142748;
   Prof_PriceDA.Data[4841] := 0.1142748;
   Prof_PriceDA.Data[4842] := 0.1142748;
   Prof_PriceDA.Data[4843] := 0.1142748;
   Prof_PriceDA.Data[4844] := 0.0986364;
   Prof_PriceDA.Data[4845] := 0.0986364;
   Prof_PriceDA.Data[4846] := 0.0986364;
   Prof_PriceDA.Data[4847] := 0.0986364;
   Prof_PriceDA.Data[4848] := 0.1005588;
   Prof_PriceDA.Data[4849] := 0.1005588;
   Prof_PriceDA.Data[4850] := 0.1005588;
   Prof_PriceDA.Data[4851] := 0.1005588;
   Prof_PriceDA.Data[4852] := 0.1060236;
   Prof_PriceDA.Data[4853] := 0.1060236;
   Prof_PriceDA.Data[4854] := 0.1060236;
   Prof_PriceDA.Data[4855] := 0.1060236;
   Prof_PriceDA.Data[4856] := 0.1154952;
   Prof_PriceDA.Data[4857] := 0.1154952;
   Prof_PriceDA.Data[4858] := 0.1154952;
   Prof_PriceDA.Data[4859] := 0.1154952;
   Prof_PriceDA.Data[4860] := 0.153846;
   Prof_PriceDA.Data[4861] := 0.153846;
   Prof_PriceDA.Data[4862] := 0.153846;
   Prof_PriceDA.Data[4863] := 0.153846;
   Prof_PriceDA.Data[4864] := 0.1964844;
   Prof_PriceDA.Data[4865] := 0.1964844;
   Prof_PriceDA.Data[4866] := 0.1964844;
   Prof_PriceDA.Data[4867] := 0.1964844;
   Prof_PriceDA.Data[4868] := 0.2781972;
   Prof_PriceDA.Data[4869] := 0.2781972;
   Prof_PriceDA.Data[4870] := 0.2781972;
   Prof_PriceDA.Data[4871] := 0.2781972;
   Prof_PriceDA.Data[4872] := 0.3032856;
   Prof_PriceDA.Data[4873] := 0.3032856;
   Prof_PriceDA.Data[4874] := 0.3032856;
   Prof_PriceDA.Data[4875] := 0.3032856;
   Prof_PriceDA.Data[4876] := 0.2709936;
   Prof_PriceDA.Data[4877] := 0.2709936;
   Prof_PriceDA.Data[4878] := 0.2709936;
   Prof_PriceDA.Data[4879] := 0.2709936;
   Prof_PriceDA.Data[4880] := 0.187596;
   Prof_PriceDA.Data[4881] := 0.187596;
   Prof_PriceDA.Data[4882] := 0.187596;
   Prof_PriceDA.Data[4883] := 0.187596;
   Prof_PriceDA.Data[4884] := 0.176904;
   Prof_PriceDA.Data[4885] := 0.176904;
   Prof_PriceDA.Data[4886] := 0.176904;
   Prof_PriceDA.Data[4887] := 0.176904;
   Prof_PriceDA.Data[4888] := 0.1739556;
   Prof_PriceDA.Data[4889] := 0.1739556;
   Prof_PriceDA.Data[4890] := 0.1739556;
   Prof_PriceDA.Data[4891] := 0.1739556;
   Prof_PriceDA.Data[4892] := 0.1439748;
   Prof_PriceDA.Data[4893] := 0.1439748;
   Prof_PriceDA.Data[4894] := 0.1439748;
   Prof_PriceDA.Data[4895] := 0.1439748;
   Prof_PriceDA.Data[4896] := 0.1269432;
   Prof_PriceDA.Data[4897] := 0.1269432;
   Prof_PriceDA.Data[4898] := 0.1269432;
   Prof_PriceDA.Data[4899] := 0.1269432;
   Prof_PriceDA.Data[4900] := 0.1223964;
   Prof_PriceDA.Data[4901] := 0.1223964;
   Prof_PriceDA.Data[4902] := 0.1223964;
   Prof_PriceDA.Data[4903] := 0.1223964;
   Prof_PriceDA.Data[4904] := 0.1204956;
   Prof_PriceDA.Data[4905] := 0.1204956;
   Prof_PriceDA.Data[4906] := 0.1204956;
   Prof_PriceDA.Data[4907] := 0.1204956;
   Prof_PriceDA.Data[4908] := 0.1224288;
   Prof_PriceDA.Data[4909] := 0.1224288;
   Prof_PriceDA.Data[4910] := 0.1224288;
   Prof_PriceDA.Data[4911] := 0.1224288;
   Prof_PriceDA.Data[4912] := 0.1231308;
   Prof_PriceDA.Data[4913] := 0.1231308;
   Prof_PriceDA.Data[4914] := 0.1231308;
   Prof_PriceDA.Data[4915] := 0.1231308;
   Prof_PriceDA.Data[4916] := 0.1458;
   Prof_PriceDA.Data[4917] := 0.1458;
   Prof_PriceDA.Data[4918] := 0.1458;
   Prof_PriceDA.Data[4919] := 0.1458;
   Prof_PriceDA.Data[4920] := 0.1756512;
   Prof_PriceDA.Data[4921] := 0.1756512;
   Prof_PriceDA.Data[4922] := 0.1756512;
   Prof_PriceDA.Data[4923] := 0.1756512;
   Prof_PriceDA.Data[4924] := 0.188244;
   Prof_PriceDA.Data[4925] := 0.188244;
   Prof_PriceDA.Data[4926] := 0.188244;
   Prof_PriceDA.Data[4927] := 0.188244;
   Prof_PriceDA.Data[4928] := 0.1582416;
   Prof_PriceDA.Data[4929] := 0.1582416;
   Prof_PriceDA.Data[4930] := 0.1582416;
   Prof_PriceDA.Data[4931] := 0.1582416;
   Prof_PriceDA.Data[4932] := 0.1398276;
   Prof_PriceDA.Data[4933] := 0.1398276;
   Prof_PriceDA.Data[4934] := 0.1398276;
   Prof_PriceDA.Data[4935] := 0.1398276;
   Prof_PriceDA.Data[4936] := 0.1123524;
   Prof_PriceDA.Data[4937] := 0.1123524;
   Prof_PriceDA.Data[4938] := 0.1123524;
   Prof_PriceDA.Data[4939] := 0.1123524;
   Prof_PriceDA.Data[4940] := 0.0950508;
   Prof_PriceDA.Data[4941] := 0.0950508;
   Prof_PriceDA.Data[4942] := 0.0950508;
   Prof_PriceDA.Data[4943] := 0.0950508;
   Prof_PriceDA.Data[4944] := 0.0867564;
   Prof_PriceDA.Data[4945] := 0.0867564;
   Prof_PriceDA.Data[4946] := 0.0867564;
   Prof_PriceDA.Data[4947] := 0.0867564;
   Prof_PriceDA.Data[4948] := 0.0860436;
   Prof_PriceDA.Data[4949] := 0.0860436;
   Prof_PriceDA.Data[4950] := 0.0860436;
   Prof_PriceDA.Data[4951] := 0.0860436;
   Prof_PriceDA.Data[4952] := 0.107892;
   Prof_PriceDA.Data[4953] := 0.107892;
   Prof_PriceDA.Data[4954] := 0.107892;
   Prof_PriceDA.Data[4955] := 0.107892;
   Prof_PriceDA.Data[4956] := 0.1171476;
   Prof_PriceDA.Data[4957] := 0.1171476;
   Prof_PriceDA.Data[4958] := 0.1171476;
   Prof_PriceDA.Data[4959] := 0.1171476;
   Prof_PriceDA.Data[4960] := 0.1718604;
   Prof_PriceDA.Data[4961] := 0.1718604;
   Prof_PriceDA.Data[4962] := 0.1718604;
   Prof_PriceDA.Data[4963] := 0.1718604;
   Prof_PriceDA.Data[4964] := 0.2034612;
   Prof_PriceDA.Data[4965] := 0.2034612;
   Prof_PriceDA.Data[4966] := 0.2034612;
   Prof_PriceDA.Data[4967] := 0.2034612;
   Prof_PriceDA.Data[4968] := 0.2067012;
   Prof_PriceDA.Data[4969] := 0.2067012;
   Prof_PriceDA.Data[4970] := 0.2067012;
   Prof_PriceDA.Data[4971] := 0.2067012;
   Prof_PriceDA.Data[4972] := 0.2070792;
   Prof_PriceDA.Data[4973] := 0.2070792;
   Prof_PriceDA.Data[4974] := 0.2070792;
   Prof_PriceDA.Data[4975] := 0.2070792;
   Prof_PriceDA.Data[4976] := 0.1797876;
   Prof_PriceDA.Data[4977] := 0.1797876;
   Prof_PriceDA.Data[4978] := 0.1797876;
   Prof_PriceDA.Data[4979] := 0.1797876;
   Prof_PriceDA.Data[4980] := 0.1654884;
   Prof_PriceDA.Data[4981] := 0.1654884;
   Prof_PriceDA.Data[4982] := 0.1654884;
   Prof_PriceDA.Data[4983] := 0.1654884;
   Prof_PriceDA.Data[4984] := 0.145422;
   Prof_PriceDA.Data[4985] := 0.145422;
   Prof_PriceDA.Data[4986] := 0.145422;
   Prof_PriceDA.Data[4987] := 0.145422;
   Prof_PriceDA.Data[4988] := 0.1260468;
   Prof_PriceDA.Data[4989] := 0.1260468;
   Prof_PriceDA.Data[4990] := 0.1260468;
   Prof_PriceDA.Data[4991] := 0.1260468;
   Prof_PriceDA.Data[4992] := 0.13203;
   Prof_PriceDA.Data[4993] := 0.13203;
   Prof_PriceDA.Data[4994] := 0.13203;
   Prof_PriceDA.Data[4995] := 0.13203;
   Prof_PriceDA.Data[4996] := 0.1259496;
   Prof_PriceDA.Data[4997] := 0.1259496;
   Prof_PriceDA.Data[4998] := 0.1259496;
   Prof_PriceDA.Data[4999] := 0.1259496;
   Prof_PriceDA.Data[5000] := 0.1227312;
   Prof_PriceDA.Data[5001] := 0.1227312;
   Prof_PriceDA.Data[5002] := 0.1227312;
   Prof_PriceDA.Data[5003] := 0.1227312;
   Prof_PriceDA.Data[5004] := 0.1168668;
   Prof_PriceDA.Data[5005] := 0.1168668;
   Prof_PriceDA.Data[5006] := 0.1168668;
   Prof_PriceDA.Data[5007] := 0.1168668;
   Prof_PriceDA.Data[5008] := 0.1191024;
   Prof_PriceDA.Data[5009] := 0.1191024;
   Prof_PriceDA.Data[5010] := 0.1191024;
   Prof_PriceDA.Data[5011] := 0.1191024;
   Prof_PriceDA.Data[5012] := 0.1260468;
   Prof_PriceDA.Data[5013] := 0.1260468;
   Prof_PriceDA.Data[5014] := 0.1260468;
   Prof_PriceDA.Data[5015] := 0.1260468;
   Prof_PriceDA.Data[5016] := 0.151794;
   Prof_PriceDA.Data[5017] := 0.151794;
   Prof_PriceDA.Data[5018] := 0.151794;
   Prof_PriceDA.Data[5019] := 0.151794;
   Prof_PriceDA.Data[5020] := 0.1414152;
   Prof_PriceDA.Data[5021] := 0.1414152;
   Prof_PriceDA.Data[5022] := 0.1414152;
   Prof_PriceDA.Data[5023] := 0.1414152;
   Prof_PriceDA.Data[5024] := 0.1065204;
   Prof_PriceDA.Data[5025] := 0.1065204;
   Prof_PriceDA.Data[5026] := 0.1065204;
   Prof_PriceDA.Data[5027] := 0.1065204;
   Prof_PriceDA.Data[5028] := 0.0763344;
   Prof_PriceDA.Data[5029] := 0.0763344;
   Prof_PriceDA.Data[5030] := 0.0763344;
   Prof_PriceDA.Data[5031] := 0.0763344;
   Prof_PriceDA.Data[5032] := 0.0634392;
   Prof_PriceDA.Data[5033] := 0.0634392;
   Prof_PriceDA.Data[5034] := 0.0634392;
   Prof_PriceDA.Data[5035] := 0.0634392;
   Prof_PriceDA.Data[5036] := 0.0612036;
   Prof_PriceDA.Data[5037] := 0.0612036;
   Prof_PriceDA.Data[5038] := 0.0612036;
   Prof_PriceDA.Data[5039] := 0.0612036;
   Prof_PriceDA.Data[5040] := 0.0569916;
   Prof_PriceDA.Data[5041] := 0.0569916;
   Prof_PriceDA.Data[5042] := 0.0569916;
   Prof_PriceDA.Data[5043] := 0.0569916;
   Prof_PriceDA.Data[5044] := 0.0606852;
   Prof_PriceDA.Data[5045] := 0.0606852;
   Prof_PriceDA.Data[5046] := 0.0606852;
   Prof_PriceDA.Data[5047] := 0.0606852;
   Prof_PriceDA.Data[5048] := 0.0737316;
   Prof_PriceDA.Data[5049] := 0.0737316;
   Prof_PriceDA.Data[5050] := 0.0737316;
   Prof_PriceDA.Data[5051] := 0.0737316;
   Prof_PriceDA.Data[5052] := 0.128358;
   Prof_PriceDA.Data[5053] := 0.128358;
   Prof_PriceDA.Data[5054] := 0.128358;
   Prof_PriceDA.Data[5055] := 0.128358;
   Prof_PriceDA.Data[5056] := 0.1802304;
   Prof_PriceDA.Data[5057] := 0.1802304;
   Prof_PriceDA.Data[5058] := 0.1802304;
   Prof_PriceDA.Data[5059] := 0.1802304;
   Prof_PriceDA.Data[5060] := 0.2145528;
   Prof_PriceDA.Data[5061] := 0.2145528;
   Prof_PriceDA.Data[5062] := 0.2145528;
   Prof_PriceDA.Data[5063] := 0.2145528;
   Prof_PriceDA.Data[5064] := 0.1995408;
   Prof_PriceDA.Data[5065] := 0.1995408;
   Prof_PriceDA.Data[5066] := 0.1995408;
   Prof_PriceDA.Data[5067] := 0.1995408;
   Prof_PriceDA.Data[5068] := 0.2117664;
   Prof_PriceDA.Data[5069] := 0.2117664;
   Prof_PriceDA.Data[5070] := 0.2117664;
   Prof_PriceDA.Data[5071] := 0.2117664;
   Prof_PriceDA.Data[5072] := 0.1919808;
   Prof_PriceDA.Data[5073] := 0.1919808;
   Prof_PriceDA.Data[5074] := 0.1919808;
   Prof_PriceDA.Data[5075] := 0.1919808;
   Prof_PriceDA.Data[5076] := 0.1703268;
   Prof_PriceDA.Data[5077] := 0.1703268;
   Prof_PriceDA.Data[5078] := 0.1703268;
   Prof_PriceDA.Data[5079] := 0.1703268;
   Prof_PriceDA.Data[5080] := 0.1657152;
   Prof_PriceDA.Data[5081] := 0.1657152;
   Prof_PriceDA.Data[5082] := 0.1657152;
   Prof_PriceDA.Data[5083] := 0.1657152;
   Prof_PriceDA.Data[5084] := 0.1615464;
   Prof_PriceDA.Data[5085] := 0.1615464;
   Prof_PriceDA.Data[5086] := 0.1615464;
   Prof_PriceDA.Data[5087] := 0.1615464;
   Prof_PriceDA.Data[5088] := 0.1378512;
   Prof_PriceDA.Data[5089] := 0.1378512;
   Prof_PriceDA.Data[5090] := 0.1378512;
   Prof_PriceDA.Data[5091] := 0.1378512;
   Prof_PriceDA.Data[5092] := 0.138294;
   Prof_PriceDA.Data[5093] := 0.138294;
   Prof_PriceDA.Data[5094] := 0.138294;
   Prof_PriceDA.Data[5095] := 0.138294;
   Prof_PriceDA.Data[5096] := 0.1283796;
   Prof_PriceDA.Data[5097] := 0.1283796;
   Prof_PriceDA.Data[5098] := 0.1283796;
   Prof_PriceDA.Data[5099] := 0.1283796;
   Prof_PriceDA.Data[5100] := 0.1277748;
   Prof_PriceDA.Data[5101] := 0.1277748;
   Prof_PriceDA.Data[5102] := 0.1277748;
   Prof_PriceDA.Data[5103] := 0.1277748;
   Prof_PriceDA.Data[5104] := 0.128736;
   Prof_PriceDA.Data[5105] := 0.128736;
   Prof_PriceDA.Data[5106] := 0.128736;
   Prof_PriceDA.Data[5107] := 0.128736;
   Prof_PriceDA.Data[5108] := 0.1349352;
   Prof_PriceDA.Data[5109] := 0.1349352;
   Prof_PriceDA.Data[5110] := 0.1349352;
   Prof_PriceDA.Data[5111] := 0.1349352;
   Prof_PriceDA.Data[5112] := 0.1454112;
   Prof_PriceDA.Data[5113] := 0.1454112;
   Prof_PriceDA.Data[5114] := 0.1454112;
   Prof_PriceDA.Data[5115] := 0.1454112;
   Prof_PriceDA.Data[5116] := 0.1423332;
   Prof_PriceDA.Data[5117] := 0.1423332;
   Prof_PriceDA.Data[5118] := 0.1423332;
   Prof_PriceDA.Data[5119] := 0.1423332;
   Prof_PriceDA.Data[5120] := 0.1270296;
   Prof_PriceDA.Data[5121] := 0.1270296;
   Prof_PriceDA.Data[5122] := 0.1270296;
   Prof_PriceDA.Data[5123] := 0.1270296;
   Prof_PriceDA.Data[5124] := 0.1109592;
   Prof_PriceDA.Data[5125] := 0.1109592;
   Prof_PriceDA.Data[5126] := 0.1109592;
   Prof_PriceDA.Data[5127] := 0.1109592;
   Prof_PriceDA.Data[5128] := 0.0945432;
   Prof_PriceDA.Data[5129] := 0.0945432;
   Prof_PriceDA.Data[5130] := 0.0945432;
   Prof_PriceDA.Data[5131] := 0.0945432;
   Prof_PriceDA.Data[5132] := 0.0962172;
   Prof_PriceDA.Data[5133] := 0.0962172;
   Prof_PriceDA.Data[5134] := 0.0962172;
   Prof_PriceDA.Data[5135] := 0.0962172;
   Prof_PriceDA.Data[5136] := 0.0814752;
   Prof_PriceDA.Data[5137] := 0.0814752;
   Prof_PriceDA.Data[5138] := 0.0814752;
   Prof_PriceDA.Data[5139] := 0.0814752;
   Prof_PriceDA.Data[5140] := 0.080838;
   Prof_PriceDA.Data[5141] := 0.080838;
   Prof_PriceDA.Data[5142] := 0.080838;
   Prof_PriceDA.Data[5143] := 0.080838;
   Prof_PriceDA.Data[5144] := 0.1136808;
   Prof_PriceDA.Data[5145] := 0.1136808;
   Prof_PriceDA.Data[5146] := 0.1136808;
   Prof_PriceDA.Data[5147] := 0.1136808;
   Prof_PriceDA.Data[5148] := 0.1515996;
   Prof_PriceDA.Data[5149] := 0.1515996;
   Prof_PriceDA.Data[5150] := 0.1515996;
   Prof_PriceDA.Data[5151] := 0.1515996;
   Prof_PriceDA.Data[5152] := 0.20547;
   Prof_PriceDA.Data[5153] := 0.20547;
   Prof_PriceDA.Data[5154] := 0.20547;
   Prof_PriceDA.Data[5155] := 0.20547;
   Prof_PriceDA.Data[5156] := 0.2142504;
   Prof_PriceDA.Data[5157] := 0.2142504;
   Prof_PriceDA.Data[5158] := 0.2142504;
   Prof_PriceDA.Data[5159] := 0.2142504;
   Prof_PriceDA.Data[5160] := 0.2108916;
   Prof_PriceDA.Data[5161] := 0.2108916;
   Prof_PriceDA.Data[5162] := 0.2108916;
   Prof_PriceDA.Data[5163] := 0.2108916;
   Prof_PriceDA.Data[5164] := 0.2121984;
   Prof_PriceDA.Data[5165] := 0.2121984;
   Prof_PriceDA.Data[5166] := 0.2121984;
   Prof_PriceDA.Data[5167] := 0.2121984;
   Prof_PriceDA.Data[5168] := 0.1816344;
   Prof_PriceDA.Data[5169] := 0.1816344;
   Prof_PriceDA.Data[5170] := 0.1816344;
   Prof_PriceDA.Data[5171] := 0.1816344;
   Prof_PriceDA.Data[5172] := 0.1752408;
   Prof_PriceDA.Data[5173] := 0.1752408;
   Prof_PriceDA.Data[5174] := 0.1752408;
   Prof_PriceDA.Data[5175] := 0.1752408;
   Prof_PriceDA.Data[5176] := 0.1579716;
   Prof_PriceDA.Data[5177] := 0.1579716;
   Prof_PriceDA.Data[5178] := 0.1579716;
   Prof_PriceDA.Data[5179] := 0.1579716;
   Prof_PriceDA.Data[5180] := 0.1437696;
   Prof_PriceDA.Data[5181] := 0.1437696;
   Prof_PriceDA.Data[5182] := 0.1437696;
   Prof_PriceDA.Data[5183] := 0.1437696;
   Prof_PriceDA.Data[5184] := 0.1412748;
   Prof_PriceDA.Data[5185] := 0.1412748;
   Prof_PriceDA.Data[5186] := 0.1412748;
   Prof_PriceDA.Data[5187] := 0.1412748;
   Prof_PriceDA.Data[5188] := 0.1266408;
   Prof_PriceDA.Data[5189] := 0.1266408;
   Prof_PriceDA.Data[5190] := 0.1266408;
   Prof_PriceDA.Data[5191] := 0.1266408;
   Prof_PriceDA.Data[5192] := 0.1217808;
   Prof_PriceDA.Data[5193] := 0.1217808;
   Prof_PriceDA.Data[5194] := 0.1217808;
   Prof_PriceDA.Data[5195] := 0.1217808;
   Prof_PriceDA.Data[5196] := 0.1202796;
   Prof_PriceDA.Data[5197] := 0.1202796;
   Prof_PriceDA.Data[5198] := 0.1202796;
   Prof_PriceDA.Data[5199] := 0.1202796;
   Prof_PriceDA.Data[5200] := 0.12393;
   Prof_PriceDA.Data[5201] := 0.12393;
   Prof_PriceDA.Data[5202] := 0.12393;
   Prof_PriceDA.Data[5203] := 0.12393;
   Prof_PriceDA.Data[5204] := 0.1646784;
   Prof_PriceDA.Data[5205] := 0.1646784;
   Prof_PriceDA.Data[5206] := 0.1646784;
   Prof_PriceDA.Data[5207] := 0.1646784;
   Prof_PriceDA.Data[5208] := 0.2244888;
   Prof_PriceDA.Data[5209] := 0.2244888;
   Prof_PriceDA.Data[5210] := 0.2244888;
   Prof_PriceDA.Data[5211] := 0.2244888;
   Prof_PriceDA.Data[5212] := 0.2619324;
   Prof_PriceDA.Data[5213] := 0.2619324;
   Prof_PriceDA.Data[5214] := 0.2619324;
   Prof_PriceDA.Data[5215] := 0.2619324;
   Prof_PriceDA.Data[5216] := 0.1898856;
   Prof_PriceDA.Data[5217] := 0.1898856;
   Prof_PriceDA.Data[5218] := 0.1898856;
   Prof_PriceDA.Data[5219] := 0.1898856;
   Prof_PriceDA.Data[5220] := 0.17928;
   Prof_PriceDA.Data[5221] := 0.17928;
   Prof_PriceDA.Data[5222] := 0.17928;
   Prof_PriceDA.Data[5223] := 0.17928;
   Prof_PriceDA.Data[5224] := 0.1571292;
   Prof_PriceDA.Data[5225] := 0.1571292;
   Prof_PriceDA.Data[5226] := 0.1571292;
   Prof_PriceDA.Data[5227] := 0.1571292;
   Prof_PriceDA.Data[5228] := 0.1439964;
   Prof_PriceDA.Data[5229] := 0.1439964;
   Prof_PriceDA.Data[5230] := 0.1439964;
   Prof_PriceDA.Data[5231] := 0.1439964;
   Prof_PriceDA.Data[5232] := 0.1381104;
   Prof_PriceDA.Data[5233] := 0.1381104;
   Prof_PriceDA.Data[5234] := 0.1381104;
   Prof_PriceDA.Data[5235] := 0.1381104;
   Prof_PriceDA.Data[5236] := 0.1377216;
   Prof_PriceDA.Data[5237] := 0.1377216;
   Prof_PriceDA.Data[5238] := 0.1377216;
   Prof_PriceDA.Data[5239] := 0.1377216;
   Prof_PriceDA.Data[5240] := 0.1576908;
   Prof_PriceDA.Data[5241] := 0.1576908;
   Prof_PriceDA.Data[5242] := 0.1576908;
   Prof_PriceDA.Data[5243] := 0.1576908;
   Prof_PriceDA.Data[5244] := 0.2053944;
   Prof_PriceDA.Data[5245] := 0.2053944;
   Prof_PriceDA.Data[5246] := 0.2053944;
   Prof_PriceDA.Data[5247] := 0.2053944;
   Prof_PriceDA.Data[5248] := 0.2542212;
   Prof_PriceDA.Data[5249] := 0.2542212;
   Prof_PriceDA.Data[5250] := 0.2542212;
   Prof_PriceDA.Data[5251] := 0.2542212;
   Prof_PriceDA.Data[5252] := 0.3007044;
   Prof_PriceDA.Data[5253] := 0.3007044;
   Prof_PriceDA.Data[5254] := 0.3007044;
   Prof_PriceDA.Data[5255] := 0.3007044;
   Prof_PriceDA.Data[5256] := 0.3385584;
   Prof_PriceDA.Data[5257] := 0.3385584;
   Prof_PriceDA.Data[5258] := 0.3385584;
   Prof_PriceDA.Data[5259] := 0.3385584;
   Prof_PriceDA.Data[5260] := 0.314172;
   Prof_PriceDA.Data[5261] := 0.314172;
   Prof_PriceDA.Data[5262] := 0.314172;
   Prof_PriceDA.Data[5263] := 0.314172;
   Prof_PriceDA.Data[5264] := 0.2235384;
   Prof_PriceDA.Data[5265] := 0.2235384;
   Prof_PriceDA.Data[5266] := 0.2235384;
   Prof_PriceDA.Data[5267] := 0.2235384;
   Prof_PriceDA.Data[5268] := 0.1914516;
   Prof_PriceDA.Data[5269] := 0.1914516;
   Prof_PriceDA.Data[5270] := 0.1914516;
   Prof_PriceDA.Data[5271] := 0.1914516;
   Prof_PriceDA.Data[5272] := 0.1759428;
   Prof_PriceDA.Data[5273] := 0.1759428;
   Prof_PriceDA.Data[5274] := 0.1759428;
   Prof_PriceDA.Data[5275] := 0.1759428;
   Prof_PriceDA.Data[5276] := 0.1442664;
   Prof_PriceDA.Data[5277] := 0.1442664;
   Prof_PriceDA.Data[5278] := 0.1442664;
   Prof_PriceDA.Data[5279] := 0.1442664;
   Prof_PriceDA.Data[5280] := 0.154332;
   Prof_PriceDA.Data[5281] := 0.154332;
   Prof_PriceDA.Data[5282] := 0.154332;
   Prof_PriceDA.Data[5283] := 0.154332;
   Prof_PriceDA.Data[5284] := 0.139428;
   Prof_PriceDA.Data[5285] := 0.139428;
   Prof_PriceDA.Data[5286] := 0.139428;
   Prof_PriceDA.Data[5287] := 0.139428;
   Prof_PriceDA.Data[5288] := 0.1344168;
   Prof_PriceDA.Data[5289] := 0.1344168;
   Prof_PriceDA.Data[5290] := 0.1344168;
   Prof_PriceDA.Data[5291] := 0.1344168;
   Prof_PriceDA.Data[5292] := 0.1337688;
   Prof_PriceDA.Data[5293] := 0.1337688;
   Prof_PriceDA.Data[5294] := 0.1337688;
   Prof_PriceDA.Data[5295] := 0.1337688;
   Prof_PriceDA.Data[5296] := 0.1378404;
   Prof_PriceDA.Data[5297] := 0.1378404;
   Prof_PriceDA.Data[5298] := 0.1378404;
   Prof_PriceDA.Data[5299] := 0.1378404;
   Prof_PriceDA.Data[5300] := 0.1590192;
   Prof_PriceDA.Data[5301] := 0.1590192;
   Prof_PriceDA.Data[5302] := 0.1590192;
   Prof_PriceDA.Data[5303] := 0.1590192;
   Prof_PriceDA.Data[5304] := 0.2322324;
   Prof_PriceDA.Data[5305] := 0.2322324;
   Prof_PriceDA.Data[5306] := 0.2322324;
   Prof_PriceDA.Data[5307] := 0.2322324;
   Prof_PriceDA.Data[5308] := 0.2833596;
   Prof_PriceDA.Data[5309] := 0.2833596;
   Prof_PriceDA.Data[5310] := 0.2833596;
   Prof_PriceDA.Data[5311] := 0.2833596;
   Prof_PriceDA.Data[5312] := 0.1877148;
   Prof_PriceDA.Data[5313] := 0.1877148;
   Prof_PriceDA.Data[5314] := 0.1877148;
   Prof_PriceDA.Data[5315] := 0.1877148;
   Prof_PriceDA.Data[5316] := 0.1683828;
   Prof_PriceDA.Data[5317] := 0.1683828;
   Prof_PriceDA.Data[5318] := 0.1683828;
   Prof_PriceDA.Data[5319] := 0.1683828;
   Prof_PriceDA.Data[5320] := 0.1544076;
   Prof_PriceDA.Data[5321] := 0.1544076;
   Prof_PriceDA.Data[5322] := 0.1544076;
   Prof_PriceDA.Data[5323] := 0.1544076;
   Prof_PriceDA.Data[5324] := 0.139374;
   Prof_PriceDA.Data[5325] := 0.139374;
   Prof_PriceDA.Data[5326] := 0.139374;
   Prof_PriceDA.Data[5327] := 0.139374;
   Prof_PriceDA.Data[5328] := 0.1379268;
   Prof_PriceDA.Data[5329] := 0.1379268;
   Prof_PriceDA.Data[5330] := 0.1379268;
   Prof_PriceDA.Data[5331] := 0.1379268;
   Prof_PriceDA.Data[5332] := 0.140346;
   Prof_PriceDA.Data[5333] := 0.140346;
   Prof_PriceDA.Data[5334] := 0.140346;
   Prof_PriceDA.Data[5335] := 0.140346;
   Prof_PriceDA.Data[5336] := 0.1505088;
   Prof_PriceDA.Data[5337] := 0.1505088;
   Prof_PriceDA.Data[5338] := 0.1505088;
   Prof_PriceDA.Data[5339] := 0.1505088;
   Prof_PriceDA.Data[5340] := 0.1666008;
   Prof_PriceDA.Data[5341] := 0.1666008;
   Prof_PriceDA.Data[5342] := 0.1666008;
   Prof_PriceDA.Data[5343] := 0.1666008;
   Prof_PriceDA.Data[5344] := 0.2288196;
   Prof_PriceDA.Data[5345] := 0.2288196;
   Prof_PriceDA.Data[5346] := 0.2288196;
   Prof_PriceDA.Data[5347] := 0.2288196;
   Prof_PriceDA.Data[5348] := 0.3069468;
   Prof_PriceDA.Data[5349] := 0.3069468;
   Prof_PriceDA.Data[5350] := 0.3069468;
   Prof_PriceDA.Data[5351] := 0.3069468;
   Prof_PriceDA.Data[5352] := 0.3333636;
   Prof_PriceDA.Data[5353] := 0.3333636;
   Prof_PriceDA.Data[5354] := 0.3333636;
   Prof_PriceDA.Data[5355] := 0.3333636;
   Prof_PriceDA.Data[5356] := 0.2880468;
   Prof_PriceDA.Data[5357] := 0.2880468;
   Prof_PriceDA.Data[5358] := 0.2880468;
   Prof_PriceDA.Data[5359] := 0.2880468;
   Prof_PriceDA.Data[5360] := 0.2162916;
   Prof_PriceDA.Data[5361] := 0.2162916;
   Prof_PriceDA.Data[5362] := 0.2162916;
   Prof_PriceDA.Data[5363] := 0.2162916;
   Prof_PriceDA.Data[5364] := 0.1727892;
   Prof_PriceDA.Data[5365] := 0.1727892;
   Prof_PriceDA.Data[5366] := 0.1727892;
   Prof_PriceDA.Data[5367] := 0.1727892;
   Prof_PriceDA.Data[5368] := 0.1578528;
   Prof_PriceDA.Data[5369] := 0.1578528;
   Prof_PriceDA.Data[5370] := 0.1578528;
   Prof_PriceDA.Data[5371] := 0.1578528;
   Prof_PriceDA.Data[5372] := 0.1416744;
   Prof_PriceDA.Data[5373] := 0.1416744;
   Prof_PriceDA.Data[5374] := 0.1416744;
   Prof_PriceDA.Data[5375] := 0.1416744;
   Prof_PriceDA.Data[5376] := 0.1348488;
   Prof_PriceDA.Data[5377] := 0.1348488;
   Prof_PriceDA.Data[5378] := 0.1348488;
   Prof_PriceDA.Data[5379] := 0.1348488;
   Prof_PriceDA.Data[5380] := 0.1326132;
   Prof_PriceDA.Data[5381] := 0.1326132;
   Prof_PriceDA.Data[5382] := 0.1326132;
   Prof_PriceDA.Data[5383] := 0.1326132;
   Prof_PriceDA.Data[5384] := 0.1286388;
   Prof_PriceDA.Data[5385] := 0.1286388;
   Prof_PriceDA.Data[5386] := 0.1286388;
   Prof_PriceDA.Data[5387] := 0.1286388;
   Prof_PriceDA.Data[5388] := 0.1282284;
   Prof_PriceDA.Data[5389] := 0.1282284;
   Prof_PriceDA.Data[5390] := 0.1282284;
   Prof_PriceDA.Data[5391] := 0.1282284;
   Prof_PriceDA.Data[5392] := 0.1286172;
   Prof_PriceDA.Data[5393] := 0.1286172;
   Prof_PriceDA.Data[5394] := 0.1286172;
   Prof_PriceDA.Data[5395] := 0.1286172;
   Prof_PriceDA.Data[5396] := 0.1369332;
   Prof_PriceDA.Data[5397] := 0.1369332;
   Prof_PriceDA.Data[5398] := 0.1369332;
   Prof_PriceDA.Data[5399] := 0.1369332;
   Prof_PriceDA.Data[5400] := 0.1886328;
   Prof_PriceDA.Data[5401] := 0.1886328;
   Prof_PriceDA.Data[5402] := 0.1886328;
   Prof_PriceDA.Data[5403] := 0.1886328;
   Prof_PriceDA.Data[5404] := 0.2148444;
   Prof_PriceDA.Data[5405] := 0.2148444;
   Prof_PriceDA.Data[5406] := 0.2148444;
   Prof_PriceDA.Data[5407] := 0.2148444;
   Prof_PriceDA.Data[5408] := 0.1917864;
   Prof_PriceDA.Data[5409] := 0.1917864;
   Prof_PriceDA.Data[5410] := 0.1917864;
   Prof_PriceDA.Data[5411] := 0.1917864;
   Prof_PriceDA.Data[5412] := 0.1698516;
   Prof_PriceDA.Data[5413] := 0.1698516;
   Prof_PriceDA.Data[5414] := 0.1698516;
   Prof_PriceDA.Data[5415] := 0.1698516;
   Prof_PriceDA.Data[5416] := 0.1571292;
   Prof_PriceDA.Data[5417] := 0.1571292;
   Prof_PriceDA.Data[5418] := 0.1571292;
   Prof_PriceDA.Data[5419] := 0.1571292;
   Prof_PriceDA.Data[5420] := 0.1430892;
   Prof_PriceDA.Data[5421] := 0.1430892;
   Prof_PriceDA.Data[5422] := 0.1430892;
   Prof_PriceDA.Data[5423] := 0.1430892;
   Prof_PriceDA.Data[5424] := 0.13122;
   Prof_PriceDA.Data[5425] := 0.13122;
   Prof_PriceDA.Data[5426] := 0.13122;
   Prof_PriceDA.Data[5427] := 0.13122;
   Prof_PriceDA.Data[5428] := 0.1323864;
   Prof_PriceDA.Data[5429] := 0.1323864;
   Prof_PriceDA.Data[5430] := 0.1323864;
   Prof_PriceDA.Data[5431] := 0.1323864;
   Prof_PriceDA.Data[5432] := 0.1405836;
   Prof_PriceDA.Data[5433] := 0.1405836;
   Prof_PriceDA.Data[5434] := 0.1405836;
   Prof_PriceDA.Data[5435] := 0.1405836;
   Prof_PriceDA.Data[5436] := 0.1608552;
   Prof_PriceDA.Data[5437] := 0.1608552;
   Prof_PriceDA.Data[5438] := 0.1608552;
   Prof_PriceDA.Data[5439] := 0.1608552;
   Prof_PriceDA.Data[5440] := 0.1918404;
   Prof_PriceDA.Data[5441] := 0.1918404;
   Prof_PriceDA.Data[5442] := 0.1918404;
   Prof_PriceDA.Data[5443] := 0.1918404;
   Prof_PriceDA.Data[5444] := 0.2159892;
   Prof_PriceDA.Data[5445] := 0.2159892;
   Prof_PriceDA.Data[5446] := 0.2159892;
   Prof_PriceDA.Data[5447] := 0.2159892;
   Prof_PriceDA.Data[5448] := 0.2162052;
   Prof_PriceDA.Data[5449] := 0.2162052;
   Prof_PriceDA.Data[5450] := 0.2162052;
   Prof_PriceDA.Data[5451] := 0.2162052;
   Prof_PriceDA.Data[5452] := 0.1993896;
   Prof_PriceDA.Data[5453] := 0.1993896;
   Prof_PriceDA.Data[5454] := 0.1993896;
   Prof_PriceDA.Data[5455] := 0.1993896;
   Prof_PriceDA.Data[5456] := 0.1851768;
   Prof_PriceDA.Data[5457] := 0.1851768;
   Prof_PriceDA.Data[5458] := 0.1851768;
   Prof_PriceDA.Data[5459] := 0.1851768;
   Prof_PriceDA.Data[5460] := 0.1579716;
   Prof_PriceDA.Data[5461] := 0.1579716;
   Prof_PriceDA.Data[5462] := 0.1579716;
   Prof_PriceDA.Data[5463] := 0.1579716;
   Prof_PriceDA.Data[5464] := 0.1453248;
   Prof_PriceDA.Data[5465] := 0.1453248;
   Prof_PriceDA.Data[5466] := 0.1453248;
   Prof_PriceDA.Data[5467] := 0.1453248;
   Prof_PriceDA.Data[5468] := 0.129816;
   Prof_PriceDA.Data[5469] := 0.129816;
   Prof_PriceDA.Data[5470] := 0.129816;
   Prof_PriceDA.Data[5471] := 0.129816;
   Prof_PriceDA.Data[5472] := 0.1205928;
   Prof_PriceDA.Data[5473] := 0.1205928;
   Prof_PriceDA.Data[5474] := 0.1205928;
   Prof_PriceDA.Data[5475] := 0.1205928;
   Prof_PriceDA.Data[5476] := 0.1121148;
   Prof_PriceDA.Data[5477] := 0.1121148;
   Prof_PriceDA.Data[5478] := 0.1121148;
   Prof_PriceDA.Data[5479] := 0.1121148;
   Prof_PriceDA.Data[5480] := 0.1109268;
   Prof_PriceDA.Data[5481] := 0.1109268;
   Prof_PriceDA.Data[5482] := 0.1109268;
   Prof_PriceDA.Data[5483] := 0.1109268;
   Prof_PriceDA.Data[5484] := 0.1096308;
   Prof_PriceDA.Data[5485] := 0.1096308;
   Prof_PriceDA.Data[5486] := 0.1096308;
   Prof_PriceDA.Data[5487] := 0.1096308;
   Prof_PriceDA.Data[5488] := 0.1096308;
   Prof_PriceDA.Data[5489] := 0.1096308;
   Prof_PriceDA.Data[5490] := 0.1096308;
   Prof_PriceDA.Data[5491] := 0.1096308;
   Prof_PriceDA.Data[5492] := 0.1193508;
   Prof_PriceDA.Data[5493] := 0.1193508;
   Prof_PriceDA.Data[5494] := 0.1193508;
   Prof_PriceDA.Data[5495] := 0.1193508;
   Prof_PriceDA.Data[5496] := 0.158328;
   Prof_PriceDA.Data[5497] := 0.158328;
   Prof_PriceDA.Data[5498] := 0.158328;
   Prof_PriceDA.Data[5499] := 0.158328;
   Prof_PriceDA.Data[5500] := 0.1742148;
   Prof_PriceDA.Data[5501] := 0.1742148;
   Prof_PriceDA.Data[5502] := 0.1742148;
   Prof_PriceDA.Data[5503] := 0.1742148;
   Prof_PriceDA.Data[5504] := 0.1794096;
   Prof_PriceDA.Data[5505] := 0.1794096;
   Prof_PriceDA.Data[5506] := 0.1794096;
   Prof_PriceDA.Data[5507] := 0.1794096;
   Prof_PriceDA.Data[5508] := 0.1623456;
   Prof_PriceDA.Data[5509] := 0.1623456;
   Prof_PriceDA.Data[5510] := 0.1623456;
   Prof_PriceDA.Data[5511] := 0.1623456;
   Prof_PriceDA.Data[5512] := 0.1463184;
   Prof_PriceDA.Data[5513] := 0.1463184;
   Prof_PriceDA.Data[5514] := 0.1463184;
   Prof_PriceDA.Data[5515] := 0.1463184;
   Prof_PriceDA.Data[5516] := 0.1380024;
   Prof_PriceDA.Data[5517] := 0.1380024;
   Prof_PriceDA.Data[5518] := 0.1380024;
   Prof_PriceDA.Data[5519] := 0.1380024;
   Prof_PriceDA.Data[5520] := 0.130626;
   Prof_PriceDA.Data[5521] := 0.130626;
   Prof_PriceDA.Data[5522] := 0.130626;
   Prof_PriceDA.Data[5523] := 0.130626;
   Prof_PriceDA.Data[5524] := 0.1261872;
   Prof_PriceDA.Data[5525] := 0.1261872;
   Prof_PriceDA.Data[5526] := 0.1261872;
   Prof_PriceDA.Data[5527] := 0.1261872;
   Prof_PriceDA.Data[5528] := 0.1297512;
   Prof_PriceDA.Data[5529] := 0.1297512;
   Prof_PriceDA.Data[5530] := 0.1297512;
   Prof_PriceDA.Data[5531] := 0.1297512;
   Prof_PriceDA.Data[5532] := 0.1470096;
   Prof_PriceDA.Data[5533] := 0.1470096;
   Prof_PriceDA.Data[5534] := 0.1470096;
   Prof_PriceDA.Data[5535] := 0.1470096;
   Prof_PriceDA.Data[5536] := 0.181764;
   Prof_PriceDA.Data[5537] := 0.181764;
   Prof_PriceDA.Data[5538] := 0.181764;
   Prof_PriceDA.Data[5539] := 0.181764;
   Prof_PriceDA.Data[5540] := 0.1843668;
   Prof_PriceDA.Data[5541] := 0.1843668;
   Prof_PriceDA.Data[5542] := 0.1843668;
   Prof_PriceDA.Data[5543] := 0.1843668;
   Prof_PriceDA.Data[5544] := 0.1918836;
   Prof_PriceDA.Data[5545] := 0.1918836;
   Prof_PriceDA.Data[5546] := 0.1918836;
   Prof_PriceDA.Data[5547] := 0.1918836;
   Prof_PriceDA.Data[5548] := 0.1853712;
   Prof_PriceDA.Data[5549] := 0.1853712;
   Prof_PriceDA.Data[5550] := 0.1853712;
   Prof_PriceDA.Data[5551] := 0.1853712;
   Prof_PriceDA.Data[5552] := 0.1789992;
   Prof_PriceDA.Data[5553] := 0.1789992;
   Prof_PriceDA.Data[5554] := 0.1789992;
   Prof_PriceDA.Data[5555] := 0.1789992;
   Prof_PriceDA.Data[5556] := 0.1529928;
   Prof_PriceDA.Data[5557] := 0.1529928;
   Prof_PriceDA.Data[5558] := 0.1529928;
   Prof_PriceDA.Data[5559] := 0.1529928;
   Prof_PriceDA.Data[5560] := 0.1429056;
   Prof_PriceDA.Data[5561] := 0.1429056;
   Prof_PriceDA.Data[5562] := 0.1429056;
   Prof_PriceDA.Data[5563] := 0.1429056;
   Prof_PriceDA.Data[5564] := 0.1239732;
   Prof_PriceDA.Data[5565] := 0.1239732;
   Prof_PriceDA.Data[5566] := 0.1239732;
   Prof_PriceDA.Data[5567] := 0.1239732;
   Prof_PriceDA.Data[5568] := 0.1306044;
   Prof_PriceDA.Data[5569] := 0.1306044;
   Prof_PriceDA.Data[5570] := 0.1306044;
   Prof_PriceDA.Data[5571] := 0.1306044;
   Prof_PriceDA.Data[5572] := 0.1193832;
   Prof_PriceDA.Data[5573] := 0.1193832;
   Prof_PriceDA.Data[5574] := 0.1193832;
   Prof_PriceDA.Data[5575] := 0.1193832;
   Prof_PriceDA.Data[5576] := 0.1181304;
   Prof_PriceDA.Data[5577] := 0.1181304;
   Prof_PriceDA.Data[5578] := 0.1181304;
   Prof_PriceDA.Data[5579] := 0.1181304;
   Prof_PriceDA.Data[5580] := 0.1156464;
   Prof_PriceDA.Data[5581] := 0.1156464;
   Prof_PriceDA.Data[5582] := 0.1156464;
   Prof_PriceDA.Data[5583] := 0.1156464;
   Prof_PriceDA.Data[5584] := 0.1216944;
   Prof_PriceDA.Data[5585] := 0.1216944;
   Prof_PriceDA.Data[5586] := 0.1216944;
   Prof_PriceDA.Data[5587] := 0.1216944;
   Prof_PriceDA.Data[5588] := 0.13392;
   Prof_PriceDA.Data[5589] := 0.13392;
   Prof_PriceDA.Data[5590] := 0.13392;
   Prof_PriceDA.Data[5591] := 0.13392;
   Prof_PriceDA.Data[5592] := 0.1674648;
   Prof_PriceDA.Data[5593] := 0.1674648;
   Prof_PriceDA.Data[5594] := 0.1674648;
   Prof_PriceDA.Data[5595] := 0.1674648;
   Prof_PriceDA.Data[5596] := 0.1978236;
   Prof_PriceDA.Data[5597] := 0.1978236;
   Prof_PriceDA.Data[5598] := 0.1978236;
   Prof_PriceDA.Data[5599] := 0.1978236;
   Prof_PriceDA.Data[5600] := 0.1741608;
   Prof_PriceDA.Data[5601] := 0.1741608;
   Prof_PriceDA.Data[5602] := 0.1741608;
   Prof_PriceDA.Data[5603] := 0.1741608;
   Prof_PriceDA.Data[5604] := 0.1593324;
   Prof_PriceDA.Data[5605] := 0.1593324;
   Prof_PriceDA.Data[5606] := 0.1593324;
   Prof_PriceDA.Data[5607] := 0.1593324;
   Prof_PriceDA.Data[5608] := 0.1399248;
   Prof_PriceDA.Data[5609] := 0.1399248;
   Prof_PriceDA.Data[5610] := 0.1399248;
   Prof_PriceDA.Data[5611] := 0.1399248;
   Prof_PriceDA.Data[5612] := 0.1272024;
   Prof_PriceDA.Data[5613] := 0.1272024;
   Prof_PriceDA.Data[5614] := 0.1272024;
   Prof_PriceDA.Data[5615] := 0.1272024;
   Prof_PriceDA.Data[5616] := 0.1191888;
   Prof_PriceDA.Data[5617] := 0.1191888;
   Prof_PriceDA.Data[5618] := 0.1191888;
   Prof_PriceDA.Data[5619] := 0.1191888;
   Prof_PriceDA.Data[5620] := 0.1188972;
   Prof_PriceDA.Data[5621] := 0.1188972;
   Prof_PriceDA.Data[5622] := 0.1188972;
   Prof_PriceDA.Data[5623] := 0.1188972;
   Prof_PriceDA.Data[5624] := 0.1216944;
   Prof_PriceDA.Data[5625] := 0.1216944;
   Prof_PriceDA.Data[5626] := 0.1216944;
   Prof_PriceDA.Data[5627] := 0.1216944;
   Prof_PriceDA.Data[5628] := 0.1370952;
   Prof_PriceDA.Data[5629] := 0.1370952;
   Prof_PriceDA.Data[5630] := 0.1370952;
   Prof_PriceDA.Data[5631] := 0.1370952;
   Prof_PriceDA.Data[5632] := 0.1721628;
   Prof_PriceDA.Data[5633] := 0.1721628;
   Prof_PriceDA.Data[5634] := 0.1721628;
   Prof_PriceDA.Data[5635] := 0.1721628;
   Prof_PriceDA.Data[5636] := 0.2049408;
   Prof_PriceDA.Data[5637] := 0.2049408;
   Prof_PriceDA.Data[5638] := 0.2049408;
   Prof_PriceDA.Data[5639] := 0.2049408;
   Prof_PriceDA.Data[5640] := 0.2110428;
   Prof_PriceDA.Data[5641] := 0.2110428;
   Prof_PriceDA.Data[5642] := 0.2110428;
   Prof_PriceDA.Data[5643] := 0.2110428;
   Prof_PriceDA.Data[5644] := 0.2149308;
   Prof_PriceDA.Data[5645] := 0.2149308;
   Prof_PriceDA.Data[5646] := 0.2149308;
   Prof_PriceDA.Data[5647] := 0.2149308;
   Prof_PriceDA.Data[5648] := 0.1967652;
   Prof_PriceDA.Data[5649] := 0.1967652;
   Prof_PriceDA.Data[5650] := 0.1967652;
   Prof_PriceDA.Data[5651] := 0.1967652;
   Prof_PriceDA.Data[5652] := 0.1700352;
   Prof_PriceDA.Data[5653] := 0.1700352;
   Prof_PriceDA.Data[5654] := 0.1700352;
   Prof_PriceDA.Data[5655] := 0.1700352;
   Prof_PriceDA.Data[5656] := 0.1497528;
   Prof_PriceDA.Data[5657] := 0.1497528;
   Prof_PriceDA.Data[5658] := 0.1497528;
   Prof_PriceDA.Data[5659] := 0.1497528;
   Prof_PriceDA.Data[5660] := 0.134946;
   Prof_PriceDA.Data[5661] := 0.134946;
   Prof_PriceDA.Data[5662] := 0.134946;
   Prof_PriceDA.Data[5663] := 0.134946;
   Prof_PriceDA.Data[5664] := 0.1395468;
   Prof_PriceDA.Data[5665] := 0.1395468;
   Prof_PriceDA.Data[5666] := 0.1395468;
   Prof_PriceDA.Data[5667] := 0.1395468;
   Prof_PriceDA.Data[5668] := 0.130464;
   Prof_PriceDA.Data[5669] := 0.130464;
   Prof_PriceDA.Data[5670] := 0.130464;
   Prof_PriceDA.Data[5671] := 0.130464;
   Prof_PriceDA.Data[5672] := 0.1266948;
   Prof_PriceDA.Data[5673] := 0.1266948;
   Prof_PriceDA.Data[5674] := 0.1266948;
   Prof_PriceDA.Data[5675] := 0.1266948;
   Prof_PriceDA.Data[5676] := 0.1222884;
   Prof_PriceDA.Data[5677] := 0.1222884;
   Prof_PriceDA.Data[5678] := 0.1222884;
   Prof_PriceDA.Data[5679] := 0.1222884;
   Prof_PriceDA.Data[5680] := 0.1193616;
   Prof_PriceDA.Data[5681] := 0.1193616;
   Prof_PriceDA.Data[5682] := 0.1193616;
   Prof_PriceDA.Data[5683] := 0.1193616;
   Prof_PriceDA.Data[5684] := 0.1248264;
   Prof_PriceDA.Data[5685] := 0.1248264;
   Prof_PriceDA.Data[5686] := 0.1248264;
   Prof_PriceDA.Data[5687] := 0.1248264;
   Prof_PriceDA.Data[5688] := 0.1381212;
   Prof_PriceDA.Data[5689] := 0.1381212;
   Prof_PriceDA.Data[5690] := 0.1381212;
   Prof_PriceDA.Data[5691] := 0.1381212;
   Prof_PriceDA.Data[5692] := 0.1493208;
   Prof_PriceDA.Data[5693] := 0.1493208;
   Prof_PriceDA.Data[5694] := 0.1493208;
   Prof_PriceDA.Data[5695] := 0.1493208;
   Prof_PriceDA.Data[5696] := 0.1511892;
   Prof_PriceDA.Data[5697] := 0.1511892;
   Prof_PriceDA.Data[5698] := 0.1511892;
   Prof_PriceDA.Data[5699] := 0.1511892;
   Prof_PriceDA.Data[5700] := 0.1508868;
   Prof_PriceDA.Data[5701] := 0.1508868;
   Prof_PriceDA.Data[5702] := 0.1508868;
   Prof_PriceDA.Data[5703] := 0.1508868;
   Prof_PriceDA.Data[5704] := 0.138024;
   Prof_PriceDA.Data[5705] := 0.138024;
   Prof_PriceDA.Data[5706] := 0.138024;
   Prof_PriceDA.Data[5707] := 0.138024;
   Prof_PriceDA.Data[5708] := 0.12393;
   Prof_PriceDA.Data[5709] := 0.12393;
   Prof_PriceDA.Data[5710] := 0.12393;
   Prof_PriceDA.Data[5711] := 0.12393;
   Prof_PriceDA.Data[5712] := 0.1121904;
   Prof_PriceDA.Data[5713] := 0.1121904;
   Prof_PriceDA.Data[5714] := 0.1121904;
   Prof_PriceDA.Data[5715] := 0.1121904;
   Prof_PriceDA.Data[5716] := 0.1080648;
   Prof_PriceDA.Data[5717] := 0.1080648;
   Prof_PriceDA.Data[5718] := 0.1080648;
   Prof_PriceDA.Data[5719] := 0.1080648;
   Prof_PriceDA.Data[5720] := 0.1125252;
   Prof_PriceDA.Data[5721] := 0.1125252;
   Prof_PriceDA.Data[5722] := 0.1125252;
   Prof_PriceDA.Data[5723] := 0.1125252;
   Prof_PriceDA.Data[5724] := 0.1363068;
   Prof_PriceDA.Data[5725] := 0.1363068;
   Prof_PriceDA.Data[5726] := 0.1363068;
   Prof_PriceDA.Data[5727] := 0.1363068;
   Prof_PriceDA.Data[5728] := 0.1677024;
   Prof_PriceDA.Data[5729] := 0.1677024;
   Prof_PriceDA.Data[5730] := 0.1677024;
   Prof_PriceDA.Data[5731] := 0.1677024;
   Prof_PriceDA.Data[5732] := 0.21735;
   Prof_PriceDA.Data[5733] := 0.21735;
   Prof_PriceDA.Data[5734] := 0.21735;
   Prof_PriceDA.Data[5735] := 0.21735;
   Prof_PriceDA.Data[5736] := 0.2160972;
   Prof_PriceDA.Data[5737] := 0.2160972;
   Prof_PriceDA.Data[5738] := 0.2160972;
   Prof_PriceDA.Data[5739] := 0.2160972;
   Prof_PriceDA.Data[5740] := 0.2048868;
   Prof_PriceDA.Data[5741] := 0.2048868;
   Prof_PriceDA.Data[5742] := 0.2048868;
   Prof_PriceDA.Data[5743] := 0.2048868;
   Prof_PriceDA.Data[5744] := 0.173556;
   Prof_PriceDA.Data[5745] := 0.173556;
   Prof_PriceDA.Data[5746] := 0.173556;
   Prof_PriceDA.Data[5747] := 0.173556;
   Prof_PriceDA.Data[5748] := 0.1505412;
   Prof_PriceDA.Data[5749] := 0.1505412;
   Prof_PriceDA.Data[5750] := 0.1505412;
   Prof_PriceDA.Data[5751] := 0.1505412;
   Prof_PriceDA.Data[5752] := 0.1351188;
   Prof_PriceDA.Data[5753] := 0.1351188;
   Prof_PriceDA.Data[5754] := 0.1351188;
   Prof_PriceDA.Data[5755] := 0.1351188;
   Prof_PriceDA.Data[5756] := 0.1295136;
   Prof_PriceDA.Data[5757] := 0.1295136;
   Prof_PriceDA.Data[5758] := 0.1295136;
   Prof_PriceDA.Data[5759] := 0.1295136;
   Prof_PriceDA.Data[5760] := 0.1363176;
   Prof_PriceDA.Data[5761] := 0.1363176;
   Prof_PriceDA.Data[5762] := 0.1363176;
   Prof_PriceDA.Data[5763] := 0.1363176;
   Prof_PriceDA.Data[5764] := 0.1292436;
   Prof_PriceDA.Data[5765] := 0.1292436;
   Prof_PriceDA.Data[5766] := 0.1292436;
   Prof_PriceDA.Data[5767] := 0.1292436;
   Prof_PriceDA.Data[5768] := 0.1137132;
   Prof_PriceDA.Data[5769] := 0.1137132;
   Prof_PriceDA.Data[5770] := 0.1137132;
   Prof_PriceDA.Data[5771] := 0.1137132;
   Prof_PriceDA.Data[5772] := 0.113724;
   Prof_PriceDA.Data[5773] := 0.113724;
   Prof_PriceDA.Data[5774] := 0.113724;
   Prof_PriceDA.Data[5775] := 0.113724;
   Prof_PriceDA.Data[5776] := 0.1215432;
   Prof_PriceDA.Data[5777] := 0.1215432;
   Prof_PriceDA.Data[5778] := 0.1215432;
   Prof_PriceDA.Data[5779] := 0.1215432;
   Prof_PriceDA.Data[5780] := 0.1246428;
   Prof_PriceDA.Data[5781] := 0.1246428;
   Prof_PriceDA.Data[5782] := 0.1246428;
   Prof_PriceDA.Data[5783] := 0.1246428;
   Prof_PriceDA.Data[5784] := 0.1444932;
   Prof_PriceDA.Data[5785] := 0.1444932;
   Prof_PriceDA.Data[5786] := 0.1444932;
   Prof_PriceDA.Data[5787] := 0.1444932;
   Prof_PriceDA.Data[5788] := 0.1420956;
   Prof_PriceDA.Data[5789] := 0.1420956;
   Prof_PriceDA.Data[5790] := 0.1420956;
   Prof_PriceDA.Data[5791] := 0.1420956;
   Prof_PriceDA.Data[5792] := 0.120906;
   Prof_PriceDA.Data[5793] := 0.120906;
   Prof_PriceDA.Data[5794] := 0.120906;
   Prof_PriceDA.Data[5795] := 0.120906;
   Prof_PriceDA.Data[5796] := 0.09612;
   Prof_PriceDA.Data[5797] := 0.09612;
   Prof_PriceDA.Data[5798] := 0.09612;
   Prof_PriceDA.Data[5799] := 0.09612;
   Prof_PriceDA.Data[5800] := 0.073764;
   Prof_PriceDA.Data[5801] := 0.073764;
   Prof_PriceDA.Data[5802] := 0.073764;
   Prof_PriceDA.Data[5803] := 0.073764;
   Prof_PriceDA.Data[5804] := 0.05292;
   Prof_PriceDA.Data[5805] := 0.05292;
   Prof_PriceDA.Data[5806] := 0.05292;
   Prof_PriceDA.Data[5807] := 0.05292;
   Prof_PriceDA.Data[5808] := 0.0297;
   Prof_PriceDA.Data[5809] := 0.0297;
   Prof_PriceDA.Data[5810] := 0.0297;
   Prof_PriceDA.Data[5811] := 0.0297;
   Prof_PriceDA.Data[5812] := 0.019008;
   Prof_PriceDA.Data[5813] := 0.019008;
   Prof_PriceDA.Data[5814] := 0.019008;
   Prof_PriceDA.Data[5815] := 0.019008;
   Prof_PriceDA.Data[5816] := 0.0572184;
   Prof_PriceDA.Data[5817] := 0.0572184;
   Prof_PriceDA.Data[5818] := 0.0572184;
   Prof_PriceDA.Data[5819] := 0.0572184;
   Prof_PriceDA.Data[5820] := 0.0780732;
   Prof_PriceDA.Data[5821] := 0.0780732;
   Prof_PriceDA.Data[5822] := 0.0780732;
   Prof_PriceDA.Data[5823] := 0.0780732;
   Prof_PriceDA.Data[5824] := 0.1435644;
   Prof_PriceDA.Data[5825] := 0.1435644;
   Prof_PriceDA.Data[5826] := 0.1435644;
   Prof_PriceDA.Data[5827] := 0.1435644;
   Prof_PriceDA.Data[5828] := 0.1693332;
   Prof_PriceDA.Data[5829] := 0.1693332;
   Prof_PriceDA.Data[5830] := 0.1693332;
   Prof_PriceDA.Data[5831] := 0.1693332;
   Prof_PriceDA.Data[5832] := 0.176526;
   Prof_PriceDA.Data[5833] := 0.176526;
   Prof_PriceDA.Data[5834] := 0.176526;
   Prof_PriceDA.Data[5835] := 0.176526;
   Prof_PriceDA.Data[5836] := 0.1771632;
   Prof_PriceDA.Data[5837] := 0.1771632;
   Prof_PriceDA.Data[5838] := 0.1771632;
   Prof_PriceDA.Data[5839] := 0.1771632;
   Prof_PriceDA.Data[5840] := 0.1706292;
   Prof_PriceDA.Data[5841] := 0.1706292;
   Prof_PriceDA.Data[5842] := 0.1706292;
   Prof_PriceDA.Data[5843] := 0.1706292;
   Prof_PriceDA.Data[5844] := 0.1626372;
   Prof_PriceDA.Data[5845] := 0.1626372;
   Prof_PriceDA.Data[5846] := 0.1626372;
   Prof_PriceDA.Data[5847] := 0.1626372;
   Prof_PriceDA.Data[5848] := 0.1358316;
   Prof_PriceDA.Data[5849] := 0.1358316;
   Prof_PriceDA.Data[5850] := 0.1358316;
   Prof_PriceDA.Data[5851] := 0.1358316;
   Prof_PriceDA.Data[5852] := 0.1227204;
   Prof_PriceDA.Data[5853] := 0.1227204;
   Prof_PriceDA.Data[5854] := 0.1227204;
   Prof_PriceDA.Data[5855] := 0.1227204;
   Prof_PriceDA.Data[5856] := 0.1238328;
   Prof_PriceDA.Data[5857] := 0.1238328;
   Prof_PriceDA.Data[5858] := 0.1238328;
   Prof_PriceDA.Data[5859] := 0.1238328;
   Prof_PriceDA.Data[5860] := 0.1172664;
   Prof_PriceDA.Data[5861] := 0.1172664;
   Prof_PriceDA.Data[5862] := 0.1172664;
   Prof_PriceDA.Data[5863] := 0.1172664;
   Prof_PriceDA.Data[5864] := 0.115668;
   Prof_PriceDA.Data[5865] := 0.115668;
   Prof_PriceDA.Data[5866] := 0.115668;
   Prof_PriceDA.Data[5867] := 0.115668;
   Prof_PriceDA.Data[5868] := 0.1113588;
   Prof_PriceDA.Data[5869] := 0.1113588;
   Prof_PriceDA.Data[5870] := 0.1113588;
   Prof_PriceDA.Data[5871] := 0.1113588;
   Prof_PriceDA.Data[5872] := 0.1151604;
   Prof_PriceDA.Data[5873] := 0.1151604;
   Prof_PriceDA.Data[5874] := 0.1151604;
   Prof_PriceDA.Data[5875] := 0.1151604;
   Prof_PriceDA.Data[5876] := 0.1288332;
   Prof_PriceDA.Data[5877] := 0.1288332;
   Prof_PriceDA.Data[5878] := 0.1288332;
   Prof_PriceDA.Data[5879] := 0.1288332;
   Prof_PriceDA.Data[5880] := 0.1513188;
   Prof_PriceDA.Data[5881] := 0.1513188;
   Prof_PriceDA.Data[5882] := 0.1513188;
   Prof_PriceDA.Data[5883] := 0.1513188;
   Prof_PriceDA.Data[5884] := 0.17604;
   Prof_PriceDA.Data[5885] := 0.17604;
   Prof_PriceDA.Data[5886] := 0.17604;
   Prof_PriceDA.Data[5887] := 0.17604;
   Prof_PriceDA.Data[5888] := 0.1595484;
   Prof_PriceDA.Data[5889] := 0.1595484;
   Prof_PriceDA.Data[5890] := 0.1595484;
   Prof_PriceDA.Data[5891] := 0.1595484;
   Prof_PriceDA.Data[5892] := 0.1176444;
   Prof_PriceDA.Data[5893] := 0.1176444;
   Prof_PriceDA.Data[5894] := 0.1176444;
   Prof_PriceDA.Data[5895] := 0.1176444;
   Prof_PriceDA.Data[5896] := 0.0878364;
   Prof_PriceDA.Data[5897] := 0.0878364;
   Prof_PriceDA.Data[5898] := 0.0878364;
   Prof_PriceDA.Data[5899] := 0.0878364;
   Prof_PriceDA.Data[5900] := 0.084618;
   Prof_PriceDA.Data[5901] := 0.084618;
   Prof_PriceDA.Data[5902] := 0.084618;
   Prof_PriceDA.Data[5903] := 0.084618;
   Prof_PriceDA.Data[5904] := 0.091476;
   Prof_PriceDA.Data[5905] := 0.091476;
   Prof_PriceDA.Data[5906] := 0.091476;
   Prof_PriceDA.Data[5907] := 0.091476;
   Prof_PriceDA.Data[5908] := 0.0626184;
   Prof_PriceDA.Data[5909] := 0.0626184;
   Prof_PriceDA.Data[5910] := 0.0626184;
   Prof_PriceDA.Data[5911] := 0.0626184;
   Prof_PriceDA.Data[5912] := 0.0921672;
   Prof_PriceDA.Data[5913] := 0.0921672;
   Prof_PriceDA.Data[5914] := 0.0921672;
   Prof_PriceDA.Data[5915] := 0.0921672;
   Prof_PriceDA.Data[5916] := 0.1216296;
   Prof_PriceDA.Data[5917] := 0.1216296;
   Prof_PriceDA.Data[5918] := 0.1216296;
   Prof_PriceDA.Data[5919] := 0.1216296;
   Prof_PriceDA.Data[5920] := 0.152766;
   Prof_PriceDA.Data[5921] := 0.152766;
   Prof_PriceDA.Data[5922] := 0.152766;
   Prof_PriceDA.Data[5923] := 0.152766;
   Prof_PriceDA.Data[5924] := 0.1925964;
   Prof_PriceDA.Data[5925] := 0.1925964;
   Prof_PriceDA.Data[5926] := 0.1925964;
   Prof_PriceDA.Data[5927] := 0.1925964;
   Prof_PriceDA.Data[5928] := 0.2588436;
   Prof_PriceDA.Data[5929] := 0.2588436;
   Prof_PriceDA.Data[5930] := 0.2588436;
   Prof_PriceDA.Data[5931] := 0.2588436;
   Prof_PriceDA.Data[5932] := 0.2024784;
   Prof_PriceDA.Data[5933] := 0.2024784;
   Prof_PriceDA.Data[5934] := 0.2024784;
   Prof_PriceDA.Data[5935] := 0.2024784;
   Prof_PriceDA.Data[5936] := 0.1784916;
   Prof_PriceDA.Data[5937] := 0.1784916;
   Prof_PriceDA.Data[5938] := 0.1784916;
   Prof_PriceDA.Data[5939] := 0.1784916;
   Prof_PriceDA.Data[5940] := 0.1745604;
   Prof_PriceDA.Data[5941] := 0.1745604;
   Prof_PriceDA.Data[5942] := 0.1745604;
   Prof_PriceDA.Data[5943] := 0.1745604;
   Prof_PriceDA.Data[5944] := 0.1605204;
   Prof_PriceDA.Data[5945] := 0.1605204;
   Prof_PriceDA.Data[5946] := 0.1605204;
   Prof_PriceDA.Data[5947] := 0.1605204;
   Prof_PriceDA.Data[5948] := 0.1555308;
   Prof_PriceDA.Data[5949] := 0.1555308;
   Prof_PriceDA.Data[5950] := 0.1555308;
   Prof_PriceDA.Data[5951] := 0.1555308;
   Prof_PriceDA.Data[5952] := 0.1387368;
   Prof_PriceDA.Data[5953] := 0.1387368;
   Prof_PriceDA.Data[5954] := 0.1387368;
   Prof_PriceDA.Data[5955] := 0.1387368;
   Prof_PriceDA.Data[5956] := 0.1302264;
   Prof_PriceDA.Data[5957] := 0.1302264;
   Prof_PriceDA.Data[5958] := 0.1302264;
   Prof_PriceDA.Data[5959] := 0.1302264;
   Prof_PriceDA.Data[5960] := 0.1188756;
   Prof_PriceDA.Data[5961] := 0.1188756;
   Prof_PriceDA.Data[5962] := 0.1188756;
   Prof_PriceDA.Data[5963] := 0.1188756;
   Prof_PriceDA.Data[5964] := 0.1167696;
   Prof_PriceDA.Data[5965] := 0.1167696;
   Prof_PriceDA.Data[5966] := 0.1167696;
   Prof_PriceDA.Data[5967] := 0.1167696;
   Prof_PriceDA.Data[5968] := 0.1265112;
   Prof_PriceDA.Data[5969] := 0.1265112;
   Prof_PriceDA.Data[5970] := 0.1265112;
   Prof_PriceDA.Data[5971] := 0.1265112;
   Prof_PriceDA.Data[5972] := 0.1686852;
   Prof_PriceDA.Data[5973] := 0.1686852;
   Prof_PriceDA.Data[5974] := 0.1686852;
   Prof_PriceDA.Data[5975] := 0.1686852;
   Prof_PriceDA.Data[5976] := 0.1939896;
   Prof_PriceDA.Data[5977] := 0.1939896;
   Prof_PriceDA.Data[5978] := 0.1939896;
   Prof_PriceDA.Data[5979] := 0.1939896;
   Prof_PriceDA.Data[5980] := 0.1906956;
   Prof_PriceDA.Data[5981] := 0.1906956;
   Prof_PriceDA.Data[5982] := 0.1906956;
   Prof_PriceDA.Data[5983] := 0.1906956;
   Prof_PriceDA.Data[5984] := 0.153306;
   Prof_PriceDA.Data[5985] := 0.153306;
   Prof_PriceDA.Data[5986] := 0.153306;
   Prof_PriceDA.Data[5987] := 0.153306;
   Prof_PriceDA.Data[5988] := 0.1248804;
   Prof_PriceDA.Data[5989] := 0.1248804;
   Prof_PriceDA.Data[5990] := 0.1248804;
   Prof_PriceDA.Data[5991] := 0.1248804;
   Prof_PriceDA.Data[5992] := 0.103302;
   Prof_PriceDA.Data[5993] := 0.103302;
   Prof_PriceDA.Data[5994] := 0.103302;
   Prof_PriceDA.Data[5995] := 0.103302;
   Prof_PriceDA.Data[5996] := 0.1115964;
   Prof_PriceDA.Data[5997] := 0.1115964;
   Prof_PriceDA.Data[5998] := 0.1115964;
   Prof_PriceDA.Data[5999] := 0.1115964;
   Prof_PriceDA.Data[6000] := 0.039798;
   Prof_PriceDA.Data[6001] := 0.039798;
   Prof_PriceDA.Data[6002] := 0.039798;
   Prof_PriceDA.Data[6003] := 0.039798;
   Prof_PriceDA.Data[6004] := 0.0315252;
   Prof_PriceDA.Data[6005] := 0.0315252;
   Prof_PriceDA.Data[6006] := 0.0315252;
   Prof_PriceDA.Data[6007] := 0.0315252;
   Prof_PriceDA.Data[6008] := 0.0721656;
   Prof_PriceDA.Data[6009] := 0.0721656;
   Prof_PriceDA.Data[6010] := 0.0721656;
   Prof_PriceDA.Data[6011] := 0.0721656;
   Prof_PriceDA.Data[6012] := 0.1109484;
   Prof_PriceDA.Data[6013] := 0.1109484;
   Prof_PriceDA.Data[6014] := 0.1109484;
   Prof_PriceDA.Data[6015] := 0.1109484;
   Prof_PriceDA.Data[6016] := 0.1677996;
   Prof_PriceDA.Data[6017] := 0.1677996;
   Prof_PriceDA.Data[6018] := 0.1677996;
   Prof_PriceDA.Data[6019] := 0.1677996;
   Prof_PriceDA.Data[6020] := 0.2093148;
   Prof_PriceDA.Data[6021] := 0.2093148;
   Prof_PriceDA.Data[6022] := 0.2093148;
   Prof_PriceDA.Data[6023] := 0.2093148;
   Prof_PriceDA.Data[6024] := 0.2734452;
   Prof_PriceDA.Data[6025] := 0.2734452;
   Prof_PriceDA.Data[6026] := 0.2734452;
   Prof_PriceDA.Data[6027] := 0.2734452;
   Prof_PriceDA.Data[6028] := 0.215298;
   Prof_PriceDA.Data[6029] := 0.215298;
   Prof_PriceDA.Data[6030] := 0.215298;
   Prof_PriceDA.Data[6031] := 0.215298;
   Prof_PriceDA.Data[6032] := 0.1860192;
   Prof_PriceDA.Data[6033] := 0.1860192;
   Prof_PriceDA.Data[6034] := 0.1860192;
   Prof_PriceDA.Data[6035] := 0.1860192;
   Prof_PriceDA.Data[6036] := 0.1675188;
   Prof_PriceDA.Data[6037] := 0.1675188;
   Prof_PriceDA.Data[6038] := 0.1675188;
   Prof_PriceDA.Data[6039] := 0.1675188;
   Prof_PriceDA.Data[6040] := 0.1552824;
   Prof_PriceDA.Data[6041] := 0.1552824;
   Prof_PriceDA.Data[6042] := 0.1552824;
   Prof_PriceDA.Data[6043] := 0.1552824;
   Prof_PriceDA.Data[6044] := 0.1442556;
   Prof_PriceDA.Data[6045] := 0.1442556;
   Prof_PriceDA.Data[6046] := 0.1442556;
   Prof_PriceDA.Data[6047] := 0.1442556;
   Prof_PriceDA.Data[6048] := 0.1448064;
   Prof_PriceDA.Data[6049] := 0.1448064;
   Prof_PriceDA.Data[6050] := 0.1448064;
   Prof_PriceDA.Data[6051] := 0.1448064;
   Prof_PriceDA.Data[6052] := 0.1312524;
   Prof_PriceDA.Data[6053] := 0.1312524;
   Prof_PriceDA.Data[6054] := 0.1312524;
   Prof_PriceDA.Data[6055] := 0.1312524;
   Prof_PriceDA.Data[6056] := 0.1238328;
   Prof_PriceDA.Data[6057] := 0.1238328;
   Prof_PriceDA.Data[6058] := 0.1238328;
   Prof_PriceDA.Data[6059] := 0.1238328;
   Prof_PriceDA.Data[6060] := 0.118854;
   Prof_PriceDA.Data[6061] := 0.118854;
   Prof_PriceDA.Data[6062] := 0.118854;
   Prof_PriceDA.Data[6063] := 0.118854;
   Prof_PriceDA.Data[6064] := 0.1313712;
   Prof_PriceDA.Data[6065] := 0.1313712;
   Prof_PriceDA.Data[6066] := 0.1313712;
   Prof_PriceDA.Data[6067] := 0.1313712;
   Prof_PriceDA.Data[6068] := 0.1473228;
   Prof_PriceDA.Data[6069] := 0.1473228;
   Prof_PriceDA.Data[6070] := 0.1473228;
   Prof_PriceDA.Data[6071] := 0.1473228;
   Prof_PriceDA.Data[6072] := 0.18387;
   Prof_PriceDA.Data[6073] := 0.18387;
   Prof_PriceDA.Data[6074] := 0.18387;
   Prof_PriceDA.Data[6075] := 0.18387;
   Prof_PriceDA.Data[6076] := 0.163944;
   Prof_PriceDA.Data[6077] := 0.163944;
   Prof_PriceDA.Data[6078] := 0.163944;
   Prof_PriceDA.Data[6079] := 0.163944;
   Prof_PriceDA.Data[6080] := 0.1172124;
   Prof_PriceDA.Data[6081] := 0.1172124;
   Prof_PriceDA.Data[6082] := 0.1172124;
   Prof_PriceDA.Data[6083] := 0.1172124;
   Prof_PriceDA.Data[6084] := 0.0805248;
   Prof_PriceDA.Data[6085] := 0.0805248;
   Prof_PriceDA.Data[6086] := 0.0805248;
   Prof_PriceDA.Data[6087] := 0.0805248;
   Prof_PriceDA.Data[6088] := 0.0244836;
   Prof_PriceDA.Data[6089] := 0.0244836;
   Prof_PriceDA.Data[6090] := 0.0244836;
   Prof_PriceDA.Data[6091] := 0.0244836;
   Prof_PriceDA.Data[6092] := 0.0119124;
   Prof_PriceDA.Data[6093] := 0.0119124;
   Prof_PriceDA.Data[6094] := 0.0119124;
   Prof_PriceDA.Data[6095] := 0.0119124;
   Prof_PriceDA.Data[6096] := 0.0075924;
   Prof_PriceDA.Data[6097] := 0.0075924;
   Prof_PriceDA.Data[6098] := 0.0075924;
   Prof_PriceDA.Data[6099] := 0.0075924;
   Prof_PriceDA.Data[6100] := 0.0011232;
   Prof_PriceDA.Data[6101] := 0.0011232;
   Prof_PriceDA.Data[6102] := 0.0011232;
   Prof_PriceDA.Data[6103] := 0.0011232;
   Prof_PriceDA.Data[6104] := 0.0041688;
   Prof_PriceDA.Data[6105] := 0.0041688;
   Prof_PriceDA.Data[6106] := 0.0041688;
   Prof_PriceDA.Data[6107] := 0.0041688;
   Prof_PriceDA.Data[6108] := 0.0786888;
   Prof_PriceDA.Data[6109] := 0.0786888;
   Prof_PriceDA.Data[6110] := 0.0786888;
   Prof_PriceDA.Data[6111] := 0.0786888;
   Prof_PriceDA.Data[6112] := 0.134892;
   Prof_PriceDA.Data[6113] := 0.134892;
   Prof_PriceDA.Data[6114] := 0.134892;
   Prof_PriceDA.Data[6115] := 0.134892;
   Prof_PriceDA.Data[6116] := 0.1743768;
   Prof_PriceDA.Data[6117] := 0.1743768;
   Prof_PriceDA.Data[6118] := 0.1743768;
   Prof_PriceDA.Data[6119] := 0.1743768;
   Prof_PriceDA.Data[6120] := 0.228744;
   Prof_PriceDA.Data[6121] := 0.228744;
   Prof_PriceDA.Data[6122] := 0.228744;
   Prof_PriceDA.Data[6123] := 0.228744;
   Prof_PriceDA.Data[6124] := 0.1930392;
   Prof_PriceDA.Data[6125] := 0.1930392;
   Prof_PriceDA.Data[6126] := 0.1930392;
   Prof_PriceDA.Data[6127] := 0.1930392;
   Prof_PriceDA.Data[6128] := 0.1734264;
   Prof_PriceDA.Data[6129] := 0.1734264;
   Prof_PriceDA.Data[6130] := 0.1734264;
   Prof_PriceDA.Data[6131] := 0.1734264;
   Prof_PriceDA.Data[6132] := 0.1610604;
   Prof_PriceDA.Data[6133] := 0.1610604;
   Prof_PriceDA.Data[6134] := 0.1610604;
   Prof_PriceDA.Data[6135] := 0.1610604;
   Prof_PriceDA.Data[6136] := 0.1397736;
   Prof_PriceDA.Data[6137] := 0.1397736;
   Prof_PriceDA.Data[6138] := 0.1397736;
   Prof_PriceDA.Data[6139] := 0.1397736;
   Prof_PriceDA.Data[6140] := 0.1315116;
   Prof_PriceDA.Data[6141] := 0.1315116;
   Prof_PriceDA.Data[6142] := 0.1315116;
   Prof_PriceDA.Data[6143] := 0.1315116;
   Prof_PriceDA.Data[6144] := 0.1128816;
   Prof_PriceDA.Data[6145] := 0.1128816;
   Prof_PriceDA.Data[6146] := 0.1128816;
   Prof_PriceDA.Data[6147] := 0.1128816;
   Prof_PriceDA.Data[6148] := 0.1133676;
   Prof_PriceDA.Data[6149] := 0.1133676;
   Prof_PriceDA.Data[6150] := 0.1133676;
   Prof_PriceDA.Data[6151] := 0.1133676;
   Prof_PriceDA.Data[6152] := 0.1125792;
   Prof_PriceDA.Data[6153] := 0.1125792;
   Prof_PriceDA.Data[6154] := 0.1125792;
   Prof_PriceDA.Data[6155] := 0.1125792;
   Prof_PriceDA.Data[6156] := 0.1146852;
   Prof_PriceDA.Data[6157] := 0.1146852;
   Prof_PriceDA.Data[6158] := 0.1146852;
   Prof_PriceDA.Data[6159] := 0.1146852;
   Prof_PriceDA.Data[6160] := 0.1219968;
   Prof_PriceDA.Data[6161] := 0.1219968;
   Prof_PriceDA.Data[6162] := 0.1219968;
   Prof_PriceDA.Data[6163] := 0.1219968;
   Prof_PriceDA.Data[6164] := 0.1468692;
   Prof_PriceDA.Data[6165] := 0.1468692;
   Prof_PriceDA.Data[6166] := 0.1468692;
   Prof_PriceDA.Data[6167] := 0.1468692;
   Prof_PriceDA.Data[6168] := 0.1857276;
   Prof_PriceDA.Data[6169] := 0.1857276;
   Prof_PriceDA.Data[6170] := 0.1857276;
   Prof_PriceDA.Data[6171] := 0.1857276;
   Prof_PriceDA.Data[6172] := 0.1662336;
   Prof_PriceDA.Data[6173] := 0.1662336;
   Prof_PriceDA.Data[6174] := 0.1662336;
   Prof_PriceDA.Data[6175] := 0.1662336;
   Prof_PriceDA.Data[6176] := 0.11718;
   Prof_PriceDA.Data[6177] := 0.11718;
   Prof_PriceDA.Data[6178] := 0.11718;
   Prof_PriceDA.Data[6179] := 0.11718;
   Prof_PriceDA.Data[6180] := 0.086076;
   Prof_PriceDA.Data[6181] := 0.086076;
   Prof_PriceDA.Data[6182] := 0.086076;
   Prof_PriceDA.Data[6183] := 0.086076;
   Prof_PriceDA.Data[6184] := 0.0622944;
   Prof_PriceDA.Data[6185] := 0.0622944;
   Prof_PriceDA.Data[6186] := 0.0622944;
   Prof_PriceDA.Data[6187] := 0.0622944;
   Prof_PriceDA.Data[6188] := 0.0057564;
   Prof_PriceDA.Data[6189] := 0.0057564;
   Prof_PriceDA.Data[6190] := 0.0057564;
   Prof_PriceDA.Data[6191] := 0.0057564;
   Prof_PriceDA.Data[6192] := 0.0016632;
   Prof_PriceDA.Data[6193] := 0.0016632;
   Prof_PriceDA.Data[6194] := 0.0016632;
   Prof_PriceDA.Data[6195] := 0.0016632;
   Prof_PriceDA.Data[6196] := 0.0007776;
   Prof_PriceDA.Data[6197] := 0.0007776;
   Prof_PriceDA.Data[6198] := 0.0007776;
   Prof_PriceDA.Data[6199] := 0.0007776;
   Prof_PriceDA.Data[6200] := 0.0142128;
   Prof_PriceDA.Data[6201] := 0.0142128;
   Prof_PriceDA.Data[6202] := 0.0142128;
   Prof_PriceDA.Data[6203] := 0.0142128;
   Prof_PriceDA.Data[6204] := 0.0805788;
   Prof_PriceDA.Data[6205] := 0.0805788;
   Prof_PriceDA.Data[6206] := 0.0805788;
   Prof_PriceDA.Data[6207] := 0.0805788;
   Prof_PriceDA.Data[6208] := 0.1324512;
   Prof_PriceDA.Data[6209] := 0.1324512;
   Prof_PriceDA.Data[6210] := 0.1324512;
   Prof_PriceDA.Data[6211] := 0.1324512;
   Prof_PriceDA.Data[6212] := 0.2071116;
   Prof_PriceDA.Data[6213] := 0.2071116;
   Prof_PriceDA.Data[6214] := 0.2071116;
   Prof_PriceDA.Data[6215] := 0.2071116;
   Prof_PriceDA.Data[6216] := 0.237006;
   Prof_PriceDA.Data[6217] := 0.237006;
   Prof_PriceDA.Data[6218] := 0.237006;
   Prof_PriceDA.Data[6219] := 0.237006;
   Prof_PriceDA.Data[6220] := 0.2223612;
   Prof_PriceDA.Data[6221] := 0.2223612;
   Prof_PriceDA.Data[6222] := 0.2223612;
   Prof_PriceDA.Data[6223] := 0.2223612;
   Prof_PriceDA.Data[6224] := 0.1900692;
   Prof_PriceDA.Data[6225] := 0.1900692;
   Prof_PriceDA.Data[6226] := 0.1900692;
   Prof_PriceDA.Data[6227] := 0.1900692;
   Prof_PriceDA.Data[6228] := 0.1577772;
   Prof_PriceDA.Data[6229] := 0.1577772;
   Prof_PriceDA.Data[6230] := 0.1577772;
   Prof_PriceDA.Data[6231] := 0.1577772;
   Prof_PriceDA.Data[6232] := 0.1492776;
   Prof_PriceDA.Data[6233] := 0.1492776;
   Prof_PriceDA.Data[6234] := 0.1492776;
   Prof_PriceDA.Data[6235] := 0.1492776;
   Prof_PriceDA.Data[6236] := 0.1302912;
   Prof_PriceDA.Data[6237] := 0.1302912;
   Prof_PriceDA.Data[6238] := 0.1302912;
   Prof_PriceDA.Data[6239] := 0.1302912;
   Prof_PriceDA.Data[6240] := 0.1153116;
   Prof_PriceDA.Data[6241] := 0.1153116;
   Prof_PriceDA.Data[6242] := 0.1153116;
   Prof_PriceDA.Data[6243] := 0.1153116;
   Prof_PriceDA.Data[6244] := 0.1140264;
   Prof_PriceDA.Data[6245] := 0.1140264;
   Prof_PriceDA.Data[6246] := 0.1140264;
   Prof_PriceDA.Data[6247] := 0.1140264;
   Prof_PriceDA.Data[6248] := 0.10854;
   Prof_PriceDA.Data[6249] := 0.10854;
   Prof_PriceDA.Data[6250] := 0.10854;
   Prof_PriceDA.Data[6251] := 0.10854;
   Prof_PriceDA.Data[6252] := 0.1099656;
   Prof_PriceDA.Data[6253] := 0.1099656;
   Prof_PriceDA.Data[6254] := 0.1099656;
   Prof_PriceDA.Data[6255] := 0.1099656;
   Prof_PriceDA.Data[6256] := 0.114048;
   Prof_PriceDA.Data[6257] := 0.114048;
   Prof_PriceDA.Data[6258] := 0.114048;
   Prof_PriceDA.Data[6259] := 0.114048;
   Prof_PriceDA.Data[6260] := 0.1347624;
   Prof_PriceDA.Data[6261] := 0.1347624;
   Prof_PriceDA.Data[6262] := 0.1347624;
   Prof_PriceDA.Data[6263] := 0.1347624;
   Prof_PriceDA.Data[6264] := 0.164322;
   Prof_PriceDA.Data[6265] := 0.164322;
   Prof_PriceDA.Data[6266] := 0.164322;
   Prof_PriceDA.Data[6267] := 0.164322;
   Prof_PriceDA.Data[6268] := 0.1642896;
   Prof_PriceDA.Data[6269] := 0.1642896;
   Prof_PriceDA.Data[6270] := 0.1642896;
   Prof_PriceDA.Data[6271] := 0.1642896;
   Prof_PriceDA.Data[6272] := 0.1339956;
   Prof_PriceDA.Data[6273] := 0.1339956;
   Prof_PriceDA.Data[6274] := 0.1339956;
   Prof_PriceDA.Data[6275] := 0.1339956;
   Prof_PriceDA.Data[6276] := 0.0899316;
   Prof_PriceDA.Data[6277] := 0.0899316;
   Prof_PriceDA.Data[6278] := 0.0899316;
   Prof_PriceDA.Data[6279] := 0.0899316;
   Prof_PriceDA.Data[6280] := 0.071064;
   Prof_PriceDA.Data[6281] := 0.071064;
   Prof_PriceDA.Data[6282] := 0.071064;
   Prof_PriceDA.Data[6283] := 0.071064;
   Prof_PriceDA.Data[6284] := 0.0343548;
   Prof_PriceDA.Data[6285] := 0.0343548;
   Prof_PriceDA.Data[6286] := 0.0343548;
   Prof_PriceDA.Data[6287] := 0.0343548;
   Prof_PriceDA.Data[6288] := 0.0138132;
   Prof_PriceDA.Data[6289] := 0.0138132;
   Prof_PriceDA.Data[6290] := 0.0138132;
   Prof_PriceDA.Data[6291] := 0.0138132;
   Prof_PriceDA.Data[6292] := 0.0086508;
   Prof_PriceDA.Data[6293] := 0.0086508;
   Prof_PriceDA.Data[6294] := 0.0086508;
   Prof_PriceDA.Data[6295] := 0.0086508;
   Prof_PriceDA.Data[6296] := 0.0415476;
   Prof_PriceDA.Data[6297] := 0.0415476;
   Prof_PriceDA.Data[6298] := 0.0415476;
   Prof_PriceDA.Data[6299] := 0.0415476;
   Prof_PriceDA.Data[6300] := 0.1037232;
   Prof_PriceDA.Data[6301] := 0.1037232;
   Prof_PriceDA.Data[6302] := 0.1037232;
   Prof_PriceDA.Data[6303] := 0.1037232;
   Prof_PriceDA.Data[6304] := 0.1464804;
   Prof_PriceDA.Data[6305] := 0.1464804;
   Prof_PriceDA.Data[6306] := 0.1464804;
   Prof_PriceDA.Data[6307] := 0.1464804;
   Prof_PriceDA.Data[6308] := 0.1729836;
   Prof_PriceDA.Data[6309] := 0.1729836;
   Prof_PriceDA.Data[6310] := 0.1729836;
   Prof_PriceDA.Data[6311] := 0.1729836;
   Prof_PriceDA.Data[6312] := 0.2413584;
   Prof_PriceDA.Data[6313] := 0.2413584;
   Prof_PriceDA.Data[6314] := 0.2413584;
   Prof_PriceDA.Data[6315] := 0.2413584;
   Prof_PriceDA.Data[6316] := 0.208764;
   Prof_PriceDA.Data[6317] := 0.208764;
   Prof_PriceDA.Data[6318] := 0.208764;
   Prof_PriceDA.Data[6319] := 0.208764;
   Prof_PriceDA.Data[6320] := 0.175068;
   Prof_PriceDA.Data[6321] := 0.175068;
   Prof_PriceDA.Data[6322] := 0.175068;
   Prof_PriceDA.Data[6323] := 0.175068;
   Prof_PriceDA.Data[6324] := 0.151524;
   Prof_PriceDA.Data[6325] := 0.151524;
   Prof_PriceDA.Data[6326] := 0.151524;
   Prof_PriceDA.Data[6327] := 0.151524;
   Prof_PriceDA.Data[6328] := 0.140994;
   Prof_PriceDA.Data[6329] := 0.140994;
   Prof_PriceDA.Data[6330] := 0.140994;
   Prof_PriceDA.Data[6331] := 0.140994;
   Prof_PriceDA.Data[6332] := 0.1352808;
   Prof_PriceDA.Data[6333] := 0.1352808;
   Prof_PriceDA.Data[6334] := 0.1352808;
   Prof_PriceDA.Data[6335] := 0.1352808;
   Prof_PriceDA.Data[6336] := 0.1441908;
   Prof_PriceDA.Data[6337] := 0.1441908;
   Prof_PriceDA.Data[6338] := 0.1441908;
   Prof_PriceDA.Data[6339] := 0.1441908;
   Prof_PriceDA.Data[6340] := 0.13662;
   Prof_PriceDA.Data[6341] := 0.13662;
   Prof_PriceDA.Data[6342] := 0.13662;
   Prof_PriceDA.Data[6343] := 0.13662;
   Prof_PriceDA.Data[6344] := 0.1405512;
   Prof_PriceDA.Data[6345] := 0.1405512;
   Prof_PriceDA.Data[6346] := 0.1405512;
   Prof_PriceDA.Data[6347] := 0.1405512;
   Prof_PriceDA.Data[6348] := 0.137808;
   Prof_PriceDA.Data[6349] := 0.137808;
   Prof_PriceDA.Data[6350] := 0.137808;
   Prof_PriceDA.Data[6351] := 0.137808;
   Prof_PriceDA.Data[6352] := 0.1404756;
   Prof_PriceDA.Data[6353] := 0.1404756;
   Prof_PriceDA.Data[6354] := 0.1404756;
   Prof_PriceDA.Data[6355] := 0.1404756;
   Prof_PriceDA.Data[6356] := 0.1484568;
   Prof_PriceDA.Data[6357] := 0.1484568;
   Prof_PriceDA.Data[6358] := 0.1484568;
   Prof_PriceDA.Data[6359] := 0.1484568;
   Prof_PriceDA.Data[6360] := 0.146016;
   Prof_PriceDA.Data[6361] := 0.146016;
   Prof_PriceDA.Data[6362] := 0.146016;
   Prof_PriceDA.Data[6363] := 0.146016;
   Prof_PriceDA.Data[6364] := 0.1347948;
   Prof_PriceDA.Data[6365] := 0.1347948;
   Prof_PriceDA.Data[6366] := 0.1347948;
   Prof_PriceDA.Data[6367] := 0.1347948;
   Prof_PriceDA.Data[6368] := 0.1058832;
   Prof_PriceDA.Data[6369] := 0.1058832;
   Prof_PriceDA.Data[6370] := 0.1058832;
   Prof_PriceDA.Data[6371] := 0.1058832;
   Prof_PriceDA.Data[6372] := 0.0783432;
   Prof_PriceDA.Data[6373] := 0.0783432;
   Prof_PriceDA.Data[6374] := 0.0783432;
   Prof_PriceDA.Data[6375] := 0.0783432;
   Prof_PriceDA.Data[6376] := 0.019494;
   Prof_PriceDA.Data[6377] := 0.019494;
   Prof_PriceDA.Data[6378] := 0.019494;
   Prof_PriceDA.Data[6379] := 0.019494;
   Prof_PriceDA.Data[6380] := 0.00243;
   Prof_PriceDA.Data[6381] := 0.00243;
   Prof_PriceDA.Data[6382] := 0.00243;
   Prof_PriceDA.Data[6383] := 0.00243;
   Prof_PriceDA.Data[6384] := 0.000864;
   Prof_PriceDA.Data[6385] := 0.000864;
   Prof_PriceDA.Data[6386] := 0.000864;
   Prof_PriceDA.Data[6387] := 0.000864;
   Prof_PriceDA.Data[6388] := 4.32E-05;
   Prof_PriceDA.Data[6389] := 4.32E-05;
   Prof_PriceDA.Data[6390] := 4.32E-05;
   Prof_PriceDA.Data[6391] := 4.32E-05;
   Prof_PriceDA.Data[6392] := 7.56E-05;
   Prof_PriceDA.Data[6393] := 7.56E-05;
   Prof_PriceDA.Data[6394] := 7.56E-05;
   Prof_PriceDA.Data[6395] := 7.56E-05;
   Prof_PriceDA.Data[6396] := 0.0650916;
   Prof_PriceDA.Data[6397] := 0.0650916;
   Prof_PriceDA.Data[6398] := 0.0650916;
   Prof_PriceDA.Data[6399] := 0.0650916;
   Prof_PriceDA.Data[6400] := 0.1236708;
   Prof_PriceDA.Data[6401] := 0.1236708;
   Prof_PriceDA.Data[6402] := 0.1236708;
   Prof_PriceDA.Data[6403] := 0.1236708;
   Prof_PriceDA.Data[6404] := 0.1769364;
   Prof_PriceDA.Data[6405] := 0.1769364;
   Prof_PriceDA.Data[6406] := 0.1769364;
   Prof_PriceDA.Data[6407] := 0.1769364;
   Prof_PriceDA.Data[6408] := 0.2254716;
   Prof_PriceDA.Data[6409] := 0.2254716;
   Prof_PriceDA.Data[6410] := 0.2254716;
   Prof_PriceDA.Data[6411] := 0.2254716;
   Prof_PriceDA.Data[6412] := 0.2034612;
   Prof_PriceDA.Data[6413] := 0.2034612;
   Prof_PriceDA.Data[6414] := 0.2034612;
   Prof_PriceDA.Data[6415] := 0.2034612;
   Prof_PriceDA.Data[6416] := 0.166914;
   Prof_PriceDA.Data[6417] := 0.166914;
   Prof_PriceDA.Data[6418] := 0.166914;
   Prof_PriceDA.Data[6419] := 0.166914;
   Prof_PriceDA.Data[6420] := 0.154116;
   Prof_PriceDA.Data[6421] := 0.154116;
   Prof_PriceDA.Data[6422] := 0.154116;
   Prof_PriceDA.Data[6423] := 0.154116;
   Prof_PriceDA.Data[6424] := 0.1454112;
   Prof_PriceDA.Data[6425] := 0.1454112;
   Prof_PriceDA.Data[6426] := 0.1454112;
   Prof_PriceDA.Data[6427] := 0.1454112;
   Prof_PriceDA.Data[6428] := 0.1249884;
   Prof_PriceDA.Data[6429] := 0.1249884;
   Prof_PriceDA.Data[6430] := 0.1249884;
   Prof_PriceDA.Data[6431] := 0.1249884;
   Prof_PriceDA.Data[6432] := 0.1188108;
   Prof_PriceDA.Data[6433] := 0.1188108;
   Prof_PriceDA.Data[6434] := 0.1188108;
   Prof_PriceDA.Data[6435] := 0.1188108;
   Prof_PriceDA.Data[6436] := 0.115452;
   Prof_PriceDA.Data[6437] := 0.115452;
   Prof_PriceDA.Data[6438] := 0.115452;
   Prof_PriceDA.Data[6439] := 0.115452;
   Prof_PriceDA.Data[6440] := 0.1132056;
   Prof_PriceDA.Data[6441] := 0.1132056;
   Prof_PriceDA.Data[6442] := 0.1132056;
   Prof_PriceDA.Data[6443] := 0.1132056;
   Prof_PriceDA.Data[6444] := 0.1155276;
   Prof_PriceDA.Data[6445] := 0.1155276;
   Prof_PriceDA.Data[6446] := 0.1155276;
   Prof_PriceDA.Data[6447] := 0.1155276;
   Prof_PriceDA.Data[6448] := 0.1188864;
   Prof_PriceDA.Data[6449] := 0.1188864;
   Prof_PriceDA.Data[6450] := 0.1188864;
   Prof_PriceDA.Data[6451] := 0.1188864;
   Prof_PriceDA.Data[6452] := 0.121716;
   Prof_PriceDA.Data[6453] := 0.121716;
   Prof_PriceDA.Data[6454] := 0.121716;
   Prof_PriceDA.Data[6455] := 0.121716;
   Prof_PriceDA.Data[6456] := 0.1188324;
   Prof_PriceDA.Data[6457] := 0.1188324;
   Prof_PriceDA.Data[6458] := 0.1188324;
   Prof_PriceDA.Data[6459] := 0.1188324;
   Prof_PriceDA.Data[6460] := 0.106218;
   Prof_PriceDA.Data[6461] := 0.106218;
   Prof_PriceDA.Data[6462] := 0.106218;
   Prof_PriceDA.Data[6463] := 0.106218;
   Prof_PriceDA.Data[6464] := 0.0736344;
   Prof_PriceDA.Data[6465] := 0.0736344;
   Prof_PriceDA.Data[6466] := 0.0736344;
   Prof_PriceDA.Data[6467] := 0.0736344;
   Prof_PriceDA.Data[6468] := 0.0316116;
   Prof_PriceDA.Data[6469] := 0.0316116;
   Prof_PriceDA.Data[6470] := 0.0316116;
   Prof_PriceDA.Data[6471] := 0.0316116;
   Prof_PriceDA.Data[6472] := 0.010908;
   Prof_PriceDA.Data[6473] := 0.010908;
   Prof_PriceDA.Data[6474] := 0.010908;
   Prof_PriceDA.Data[6475] := 0.010908;
   Prof_PriceDA.Data[6476] := 0.0016416;
   Prof_PriceDA.Data[6477] := 0.0016416;
   Prof_PriceDA.Data[6478] := 0.0016416;
   Prof_PriceDA.Data[6479] := 0.0016416;
   Prof_PriceDA.Data[6480] := 0.000702;
   Prof_PriceDA.Data[6481] := 0.000702;
   Prof_PriceDA.Data[6482] := 0.000702;
   Prof_PriceDA.Data[6483] := 0.000702;
   Prof_PriceDA.Data[6484] := -0.0003456;
   Prof_PriceDA.Data[6485] := -0.0003456;
   Prof_PriceDA.Data[6486] := -0.0003456;
   Prof_PriceDA.Data[6487] := -0.0003456;
   Prof_PriceDA.Data[6488] := 0.0007884;
   Prof_PriceDA.Data[6489] := 0.0007884;
   Prof_PriceDA.Data[6490] := 0.0007884;
   Prof_PriceDA.Data[6491] := 0.0007884;
   Prof_PriceDA.Data[6492] := 0.0187812;
   Prof_PriceDA.Data[6493] := 0.0187812;
   Prof_PriceDA.Data[6494] := 0.0187812;
   Prof_PriceDA.Data[6495] := 0.0187812;
   Prof_PriceDA.Data[6496] := 0.1079352;
   Prof_PriceDA.Data[6497] := 0.1079352;
   Prof_PriceDA.Data[6498] := 0.1079352;
   Prof_PriceDA.Data[6499] := 0.1079352;
   Prof_PriceDA.Data[6500] := 0.149796;
   Prof_PriceDA.Data[6501] := 0.149796;
   Prof_PriceDA.Data[6502] := 0.149796;
   Prof_PriceDA.Data[6503] := 0.149796;
   Prof_PriceDA.Data[6504] := 0.1598832;
   Prof_PriceDA.Data[6505] := 0.1598832;
   Prof_PriceDA.Data[6506] := 0.1598832;
   Prof_PriceDA.Data[6507] := 0.1598832;
   Prof_PriceDA.Data[6508] := 0.158166;
   Prof_PriceDA.Data[6509] := 0.158166;
   Prof_PriceDA.Data[6510] := 0.158166;
   Prof_PriceDA.Data[6511] := 0.158166;
   Prof_PriceDA.Data[6512] := 0.148824;
   Prof_PriceDA.Data[6513] := 0.148824;
   Prof_PriceDA.Data[6514] := 0.148824;
   Prof_PriceDA.Data[6515] := 0.148824;
   Prof_PriceDA.Data[6516] := 0.1400328;
   Prof_PriceDA.Data[6517] := 0.1400328;
   Prof_PriceDA.Data[6518] := 0.1400328;
   Prof_PriceDA.Data[6519] := 0.1400328;
   Prof_PriceDA.Data[6520] := 0.125334;
   Prof_PriceDA.Data[6521] := 0.125334;
   Prof_PriceDA.Data[6522] := 0.125334;
   Prof_PriceDA.Data[6523] := 0.125334;
   Prof_PriceDA.Data[6524] := 0.119502;
   Prof_PriceDA.Data[6525] := 0.119502;
   Prof_PriceDA.Data[6526] := 0.119502;
   Prof_PriceDA.Data[6527] := 0.119502;
   Prof_PriceDA.Data[6528] := 0.10692;
   Prof_PriceDA.Data[6529] := 0.10692;
   Prof_PriceDA.Data[6530] := 0.10692;
   Prof_PriceDA.Data[6531] := 0.10692;
   Prof_PriceDA.Data[6532] := 0.105948;
   Prof_PriceDA.Data[6533] := 0.105948;
   Prof_PriceDA.Data[6534] := 0.105948;
   Prof_PriceDA.Data[6535] := 0.105948;
   Prof_PriceDA.Data[6536] := 0.1073304;
   Prof_PriceDA.Data[6537] := 0.1073304;
   Prof_PriceDA.Data[6538] := 0.1073304;
   Prof_PriceDA.Data[6539] := 0.1073304;
   Prof_PriceDA.Data[6540] := 0.1075032;
   Prof_PriceDA.Data[6541] := 0.1075032;
   Prof_PriceDA.Data[6542] := 0.1075032;
   Prof_PriceDA.Data[6543] := 0.1075032;
   Prof_PriceDA.Data[6544] := 0.107838;
   Prof_PriceDA.Data[6545] := 0.107838;
   Prof_PriceDA.Data[6546] := 0.107838;
   Prof_PriceDA.Data[6547] := 0.107838;
   Prof_PriceDA.Data[6548] := 0.1214136;
   Prof_PriceDA.Data[6549] := 0.1214136;
   Prof_PriceDA.Data[6550] := 0.1214136;
   Prof_PriceDA.Data[6551] := 0.1214136;
   Prof_PriceDA.Data[6552] := 0.1614492;
   Prof_PriceDA.Data[6553] := 0.1614492;
   Prof_PriceDA.Data[6554] := 0.1614492;
   Prof_PriceDA.Data[6555] := 0.1614492;
   Prof_PriceDA.Data[6556] := 0.1707372;
   Prof_PriceDA.Data[6557] := 0.1707372;
   Prof_PriceDA.Data[6558] := 0.1707372;
   Prof_PriceDA.Data[6559] := 0.1707372;
   Prof_PriceDA.Data[6560] := 0.144612;
   Prof_PriceDA.Data[6561] := 0.144612;
   Prof_PriceDA.Data[6562] := 0.144612;
   Prof_PriceDA.Data[6563] := 0.144612;
   Prof_PriceDA.Data[6564] := 0.1070604;
   Prof_PriceDA.Data[6565] := 0.1070604;
   Prof_PriceDA.Data[6566] := 0.1070604;
   Prof_PriceDA.Data[6567] := 0.1070604;
   Prof_PriceDA.Data[6568] := 0.0843588;
   Prof_PriceDA.Data[6569] := 0.0843588;
   Prof_PriceDA.Data[6570] := 0.0843588;
   Prof_PriceDA.Data[6571] := 0.0843588;
   Prof_PriceDA.Data[6572] := 0.0798876;
   Prof_PriceDA.Data[6573] := 0.0798876;
   Prof_PriceDA.Data[6574] := 0.0798876;
   Prof_PriceDA.Data[6575] := 0.0798876;
   Prof_PriceDA.Data[6576] := 0.0821016;
   Prof_PriceDA.Data[6577] := 0.0821016;
   Prof_PriceDA.Data[6578] := 0.0821016;
   Prof_PriceDA.Data[6579] := 0.0821016;
   Prof_PriceDA.Data[6580] := 0.0835056;
   Prof_PriceDA.Data[6581] := 0.0835056;
   Prof_PriceDA.Data[6582] := 0.0835056;
   Prof_PriceDA.Data[6583] := 0.0835056;
   Prof_PriceDA.Data[6584] := 0.0917568;
   Prof_PriceDA.Data[6585] := 0.0917568;
   Prof_PriceDA.Data[6586] := 0.0917568;
   Prof_PriceDA.Data[6587] := 0.0917568;
   Prof_PriceDA.Data[6588] := 0.1085508;
   Prof_PriceDA.Data[6589] := 0.1085508;
   Prof_PriceDA.Data[6590] := 0.1085508;
   Prof_PriceDA.Data[6591] := 0.1085508;
   Prof_PriceDA.Data[6592] := 0.1429704;
   Prof_PriceDA.Data[6593] := 0.1429704;
   Prof_PriceDA.Data[6594] := 0.1429704;
   Prof_PriceDA.Data[6595] := 0.1429704;
   Prof_PriceDA.Data[6596] := 0.1568592;
   Prof_PriceDA.Data[6597] := 0.1568592;
   Prof_PriceDA.Data[6598] := 0.1568592;
   Prof_PriceDA.Data[6599] := 0.1568592;
   Prof_PriceDA.Data[6600] := 0.1869804;
   Prof_PriceDA.Data[6601] := 0.1869804;
   Prof_PriceDA.Data[6602] := 0.1869804;
   Prof_PriceDA.Data[6603] := 0.1869804;
   Prof_PriceDA.Data[6604] := 0.171828;
   Prof_PriceDA.Data[6605] := 0.171828;
   Prof_PriceDA.Data[6606] := 0.171828;
   Prof_PriceDA.Data[6607] := 0.171828;
   Prof_PriceDA.Data[6608] := 0.1521828;
   Prof_PriceDA.Data[6609] := 0.1521828;
   Prof_PriceDA.Data[6610] := 0.1521828;
   Prof_PriceDA.Data[6611] := 0.1521828;
   Prof_PriceDA.Data[6612] := 0.1384992;
   Prof_PriceDA.Data[6613] := 0.1384992;
   Prof_PriceDA.Data[6614] := 0.1384992;
   Prof_PriceDA.Data[6615] := 0.1384992;
   Prof_PriceDA.Data[6616] := 0.1163376;
   Prof_PriceDA.Data[6617] := 0.1163376;
   Prof_PriceDA.Data[6618] := 0.1163376;
   Prof_PriceDA.Data[6619] := 0.1163376;
   Prof_PriceDA.Data[6620] := 0.1065528;
   Prof_PriceDA.Data[6621] := 0.1065528;
   Prof_PriceDA.Data[6622] := 0.1065528;
   Prof_PriceDA.Data[6623] := 0.1065528;
   Prof_PriceDA.Data[6624] := 0.114426;
   Prof_PriceDA.Data[6625] := 0.114426;
   Prof_PriceDA.Data[6626] := 0.114426;
   Prof_PriceDA.Data[6627] := 0.114426;
   Prof_PriceDA.Data[6628] := 0.1117476;
   Prof_PriceDA.Data[6629] := 0.1117476;
   Prof_PriceDA.Data[6630] := 0.1117476;
   Prof_PriceDA.Data[6631] := 0.1117476;
   Prof_PriceDA.Data[6632] := 0.1086804;
   Prof_PriceDA.Data[6633] := 0.1086804;
   Prof_PriceDA.Data[6634] := 0.1086804;
   Prof_PriceDA.Data[6635] := 0.1086804;
   Prof_PriceDA.Data[6636] := 0.1099332;
   Prof_PriceDA.Data[6637] := 0.1099332;
   Prof_PriceDA.Data[6638] := 0.1099332;
   Prof_PriceDA.Data[6639] := 0.1099332;
   Prof_PriceDA.Data[6640] := 0.1132272;
   Prof_PriceDA.Data[6641] := 0.1132272;
   Prof_PriceDA.Data[6642] := 0.1132272;
   Prof_PriceDA.Data[6643] := 0.1132272;
   Prof_PriceDA.Data[6644] := 0.1220832;
   Prof_PriceDA.Data[6645] := 0.1220832;
   Prof_PriceDA.Data[6646] := 0.1220832;
   Prof_PriceDA.Data[6647] := 0.1220832;
   Prof_PriceDA.Data[6648] := 0.1521828;
   Prof_PriceDA.Data[6649] := 0.1521828;
   Prof_PriceDA.Data[6650] := 0.1521828;
   Prof_PriceDA.Data[6651] := 0.1521828;
   Prof_PriceDA.Data[6652] := 0.1583064;
   Prof_PriceDA.Data[6653] := 0.1583064;
   Prof_PriceDA.Data[6654] := 0.1583064;
   Prof_PriceDA.Data[6655] := 0.1583064;
   Prof_PriceDA.Data[6656] := 0.1551744;
   Prof_PriceDA.Data[6657] := 0.1551744;
   Prof_PriceDA.Data[6658] := 0.1551744;
   Prof_PriceDA.Data[6659] := 0.1551744;
   Prof_PriceDA.Data[6660] := 0.1403568;
   Prof_PriceDA.Data[6661] := 0.1403568;
   Prof_PriceDA.Data[6662] := 0.1403568;
   Prof_PriceDA.Data[6663] := 0.1403568;
   Prof_PriceDA.Data[6664] := 0.1103544;
   Prof_PriceDA.Data[6665] := 0.1103544;
   Prof_PriceDA.Data[6666] := 0.1103544;
   Prof_PriceDA.Data[6667] := 0.1103544;
   Prof_PriceDA.Data[6668] := 0.1058724;
   Prof_PriceDA.Data[6669] := 0.1058724;
   Prof_PriceDA.Data[6670] := 0.1058724;
   Prof_PriceDA.Data[6671] := 0.1058724;
   Prof_PriceDA.Data[6672] := 0.1052568;
   Prof_PriceDA.Data[6673] := 0.1052568;
   Prof_PriceDA.Data[6674] := 0.1052568;
   Prof_PriceDA.Data[6675] := 0.1052568;
   Prof_PriceDA.Data[6676] := 0.1080432;
   Prof_PriceDA.Data[6677] := 0.1080432;
   Prof_PriceDA.Data[6678] := 0.1080432;
   Prof_PriceDA.Data[6679] := 0.1080432;
   Prof_PriceDA.Data[6680] := 0.1128168;
   Prof_PriceDA.Data[6681] := 0.1128168;
   Prof_PriceDA.Data[6682] := 0.1128168;
   Prof_PriceDA.Data[6683] := 0.1128168;
   Prof_PriceDA.Data[6684] := 0.1251504;
   Prof_PriceDA.Data[6685] := 0.1251504;
   Prof_PriceDA.Data[6686] := 0.1251504;
   Prof_PriceDA.Data[6687] := 0.1251504;
   Prof_PriceDA.Data[6688] := 0.1503792;
   Prof_PriceDA.Data[6689] := 0.1503792;
   Prof_PriceDA.Data[6690] := 0.1503792;
   Prof_PriceDA.Data[6691] := 0.1503792;
   Prof_PriceDA.Data[6692] := 0.1712016;
   Prof_PriceDA.Data[6693] := 0.1712016;
   Prof_PriceDA.Data[6694] := 0.1712016;
   Prof_PriceDA.Data[6695] := 0.1712016;
   Prof_PriceDA.Data[6696] := 0.205632;
   Prof_PriceDA.Data[6697] := 0.205632;
   Prof_PriceDA.Data[6698] := 0.205632;
   Prof_PriceDA.Data[6699] := 0.205632;
   Prof_PriceDA.Data[6700] := 0.1912248;
   Prof_PriceDA.Data[6701] := 0.1912248;
   Prof_PriceDA.Data[6702] := 0.1912248;
   Prof_PriceDA.Data[6703] := 0.1912248;
   Prof_PriceDA.Data[6704] := 0.1594512;
   Prof_PriceDA.Data[6705] := 0.1594512;
   Prof_PriceDA.Data[6706] := 0.1594512;
   Prof_PriceDA.Data[6707] := 0.1594512;
   Prof_PriceDA.Data[6708] := 0.1449036;
   Prof_PriceDA.Data[6709] := 0.1449036;
   Prof_PriceDA.Data[6710] := 0.1449036;
   Prof_PriceDA.Data[6711] := 0.1449036;
   Prof_PriceDA.Data[6712] := 0.1326996;
   Prof_PriceDA.Data[6713] := 0.1326996;
   Prof_PriceDA.Data[6714] := 0.1326996;
   Prof_PriceDA.Data[6715] := 0.1326996;
   Prof_PriceDA.Data[6716] := 0.1161864;
   Prof_PriceDA.Data[6717] := 0.1161864;
   Prof_PriceDA.Data[6718] := 0.1161864;
   Prof_PriceDA.Data[6719] := 0.1161864;
   Prof_PriceDA.Data[6720] := 0.1102356;
   Prof_PriceDA.Data[6721] := 0.1102356;
   Prof_PriceDA.Data[6722] := 0.1102356;
   Prof_PriceDA.Data[6723] := 0.1102356;
   Prof_PriceDA.Data[6724] := 0.1087776;
   Prof_PriceDA.Data[6725] := 0.1087776;
   Prof_PriceDA.Data[6726] := 0.1087776;
   Prof_PriceDA.Data[6727] := 0.1087776;
   Prof_PriceDA.Data[6728] := 0.1059912;
   Prof_PriceDA.Data[6729] := 0.1059912;
   Prof_PriceDA.Data[6730] := 0.1059912;
   Prof_PriceDA.Data[6731] := 0.1059912;
   Prof_PriceDA.Data[6732] := 0.1063044;
   Prof_PriceDA.Data[6733] := 0.1063044;
   Prof_PriceDA.Data[6734] := 0.1063044;
   Prof_PriceDA.Data[6735] := 0.1063044;
   Prof_PriceDA.Data[6736] := 0.1118664;
   Prof_PriceDA.Data[6737] := 0.1118664;
   Prof_PriceDA.Data[6738] := 0.1118664;
   Prof_PriceDA.Data[6739] := 0.1118664;
   Prof_PriceDA.Data[6740] := 0.122418;
   Prof_PriceDA.Data[6741] := 0.122418;
   Prof_PriceDA.Data[6742] := 0.122418;
   Prof_PriceDA.Data[6743] := 0.122418;
   Prof_PriceDA.Data[6744] := 0.1487052;
   Prof_PriceDA.Data[6745] := 0.1487052;
   Prof_PriceDA.Data[6746] := 0.1487052;
   Prof_PriceDA.Data[6747] := 0.1487052;
   Prof_PriceDA.Data[6748] := 0.1657152;
   Prof_PriceDA.Data[6749] := 0.1657152;
   Prof_PriceDA.Data[6750] := 0.1657152;
   Prof_PriceDA.Data[6751] := 0.1657152;
   Prof_PriceDA.Data[6752] := 0.1566972;
   Prof_PriceDA.Data[6753] := 0.1566972;
   Prof_PriceDA.Data[6754] := 0.1566972;
   Prof_PriceDA.Data[6755] := 0.1566972;
   Prof_PriceDA.Data[6756] := 0.135;
   Prof_PriceDA.Data[6757] := 0.135;
   Prof_PriceDA.Data[6758] := 0.135;
   Prof_PriceDA.Data[6759] := 0.135;
   Prof_PriceDA.Data[6760] := 0.110376;
   Prof_PriceDA.Data[6761] := 0.110376;
   Prof_PriceDA.Data[6762] := 0.110376;
   Prof_PriceDA.Data[6763] := 0.110376;
   Prof_PriceDA.Data[6764] := 0.1075248;
   Prof_PriceDA.Data[6765] := 0.1075248;
   Prof_PriceDA.Data[6766] := 0.1075248;
   Prof_PriceDA.Data[6767] := 0.1075248;
   Prof_PriceDA.Data[6768] := 0.1059048;
   Prof_PriceDA.Data[6769] := 0.1059048;
   Prof_PriceDA.Data[6770] := 0.1059048;
   Prof_PriceDA.Data[6771] := 0.1059048;
   Prof_PriceDA.Data[6772] := 0.1074924;
   Prof_PriceDA.Data[6773] := 0.1074924;
   Prof_PriceDA.Data[6774] := 0.1074924;
   Prof_PriceDA.Data[6775] := 0.1074924;
   Prof_PriceDA.Data[6776] := 0.1098576;
   Prof_PriceDA.Data[6777] := 0.1098576;
   Prof_PriceDA.Data[6778] := 0.1098576;
   Prof_PriceDA.Data[6779] := 0.1098576;
   Prof_PriceDA.Data[6780] := 0.1288764;
   Prof_PriceDA.Data[6781] := 0.1288764;
   Prof_PriceDA.Data[6782] := 0.1288764;
   Prof_PriceDA.Data[6783] := 0.1288764;
   Prof_PriceDA.Data[6784] := 0.1465776;
   Prof_PriceDA.Data[6785] := 0.1465776;
   Prof_PriceDA.Data[6786] := 0.1465776;
   Prof_PriceDA.Data[6787] := 0.1465776;
   Prof_PriceDA.Data[6788] := 0.1611252;
   Prof_PriceDA.Data[6789] := 0.1611252;
   Prof_PriceDA.Data[6790] := 0.1611252;
   Prof_PriceDA.Data[6791] := 0.1611252;
   Prof_PriceDA.Data[6792] := 0.205578;
   Prof_PriceDA.Data[6793] := 0.205578;
   Prof_PriceDA.Data[6794] := 0.205578;
   Prof_PriceDA.Data[6795] := 0.205578;
   Prof_PriceDA.Data[6796] := 0.1930068;
   Prof_PriceDA.Data[6797] := 0.1930068;
   Prof_PriceDA.Data[6798] := 0.1930068;
   Prof_PriceDA.Data[6799] := 0.1930068;
   Prof_PriceDA.Data[6800] := 0.1576692;
   Prof_PriceDA.Data[6801] := 0.1576692;
   Prof_PriceDA.Data[6802] := 0.1576692;
   Prof_PriceDA.Data[6803] := 0.1576692;
   Prof_PriceDA.Data[6804] := 0.142776;
   Prof_PriceDA.Data[6805] := 0.142776;
   Prof_PriceDA.Data[6806] := 0.142776;
   Prof_PriceDA.Data[6807] := 0.142776;
   Prof_PriceDA.Data[6808] := 0.1296;
   Prof_PriceDA.Data[6809] := 0.1296;
   Prof_PriceDA.Data[6810] := 0.1296;
   Prof_PriceDA.Data[6811] := 0.1296;
   Prof_PriceDA.Data[6812] := 0.1187028;
   Prof_PriceDA.Data[6813] := 0.1187028;
   Prof_PriceDA.Data[6814] := 0.1187028;
   Prof_PriceDA.Data[6815] := 0.1187028;
   Prof_PriceDA.Data[6816] := 0.1152576;
   Prof_PriceDA.Data[6817] := 0.1152576;
   Prof_PriceDA.Data[6818] := 0.1152576;
   Prof_PriceDA.Data[6819] := 0.1152576;
   Prof_PriceDA.Data[6820] := 0.0640764;
   Prof_PriceDA.Data[6821] := 0.0640764;
   Prof_PriceDA.Data[6822] := 0.0640764;
   Prof_PriceDA.Data[6823] := 0.0640764;
   Prof_PriceDA.Data[6824] := 0.0236844;
   Prof_PriceDA.Data[6825] := 0.0236844;
   Prof_PriceDA.Data[6826] := 0.0236844;
   Prof_PriceDA.Data[6827] := 0.0236844;
   Prof_PriceDA.Data[6828] := 0.0324216;
   Prof_PriceDA.Data[6829] := 0.0324216;
   Prof_PriceDA.Data[6830] := 0.0324216;
   Prof_PriceDA.Data[6831] := 0.0324216;
   Prof_PriceDA.Data[6832] := 0.0692064;
   Prof_PriceDA.Data[6833] := 0.0692064;
   Prof_PriceDA.Data[6834] := 0.0692064;
   Prof_PriceDA.Data[6835] := 0.0692064;
   Prof_PriceDA.Data[6836] := 0.1137564;
   Prof_PriceDA.Data[6837] := 0.1137564;
   Prof_PriceDA.Data[6838] := 0.1137564;
   Prof_PriceDA.Data[6839] := 0.1137564;
   Prof_PriceDA.Data[6840] := 0.1436292;
   Prof_PriceDA.Data[6841] := 0.1436292;
   Prof_PriceDA.Data[6842] := 0.1436292;
   Prof_PriceDA.Data[6843] := 0.1436292;
   Prof_PriceDA.Data[6844] := 0.1567836;
   Prof_PriceDA.Data[6845] := 0.1567836;
   Prof_PriceDA.Data[6846] := 0.1567836;
   Prof_PriceDA.Data[6847] := 0.1567836;
   Prof_PriceDA.Data[6848] := 0.141912;
   Prof_PriceDA.Data[6849] := 0.141912;
   Prof_PriceDA.Data[6850] := 0.141912;
   Prof_PriceDA.Data[6851] := 0.141912;
   Prof_PriceDA.Data[6852] := 0.1055592;
   Prof_PriceDA.Data[6853] := 0.1055592;
   Prof_PriceDA.Data[6854] := 0.1055592;
   Prof_PriceDA.Data[6855] := 0.1055592;
   Prof_PriceDA.Data[6856] := 0.1039932;
   Prof_PriceDA.Data[6857] := 0.1039932;
   Prof_PriceDA.Data[6858] := 0.1039932;
   Prof_PriceDA.Data[6859] := 0.1039932;
   Prof_PriceDA.Data[6860] := 0.0934092;
   Prof_PriceDA.Data[6861] := 0.0934092;
   Prof_PriceDA.Data[6862] := 0.0934092;
   Prof_PriceDA.Data[6863] := 0.0934092;
   Prof_PriceDA.Data[6864] := 0.0904392;
   Prof_PriceDA.Data[6865] := 0.0904392;
   Prof_PriceDA.Data[6866] := 0.0904392;
   Prof_PriceDA.Data[6867] := 0.0904392;
   Prof_PriceDA.Data[6868] := 0.0753192;
   Prof_PriceDA.Data[6869] := 0.0753192;
   Prof_PriceDA.Data[6870] := 0.0753192;
   Prof_PriceDA.Data[6871] := 0.0753192;
   Prof_PriceDA.Data[6872] := 0.094176;
   Prof_PriceDA.Data[6873] := 0.094176;
   Prof_PriceDA.Data[6874] := 0.094176;
   Prof_PriceDA.Data[6875] := 0.094176;
   Prof_PriceDA.Data[6876] := 0.11664;
   Prof_PriceDA.Data[6877] := 0.11664;
   Prof_PriceDA.Data[6878] := 0.11664;
   Prof_PriceDA.Data[6879] := 0.11664;
   Prof_PriceDA.Data[6880] := 0.1324296;
   Prof_PriceDA.Data[6881] := 0.1324296;
   Prof_PriceDA.Data[6882] := 0.1324296;
   Prof_PriceDA.Data[6883] := 0.1324296;
   Prof_PriceDA.Data[6884] := 0.1532628;
   Prof_PriceDA.Data[6885] := 0.1532628;
   Prof_PriceDA.Data[6886] := 0.1532628;
   Prof_PriceDA.Data[6887] := 0.1532628;
   Prof_PriceDA.Data[6888] := 0.179334;
   Prof_PriceDA.Data[6889] := 0.179334;
   Prof_PriceDA.Data[6890] := 0.179334;
   Prof_PriceDA.Data[6891] := 0.179334;
   Prof_PriceDA.Data[6892] := 0.1873476;
   Prof_PriceDA.Data[6893] := 0.1873476;
   Prof_PriceDA.Data[6894] := 0.1873476;
   Prof_PriceDA.Data[6895] := 0.1873476;
   Prof_PriceDA.Data[6896] := 0.16092;
   Prof_PriceDA.Data[6897] := 0.16092;
   Prof_PriceDA.Data[6898] := 0.16092;
   Prof_PriceDA.Data[6899] := 0.16092;
   Prof_PriceDA.Data[6900] := 0.1465452;
   Prof_PriceDA.Data[6901] := 0.1465452;
   Prof_PriceDA.Data[6902] := 0.1465452;
   Prof_PriceDA.Data[6903] := 0.1465452;
   Prof_PriceDA.Data[6904] := 0.1107216;
   Prof_PriceDA.Data[6905] := 0.1107216;
   Prof_PriceDA.Data[6906] := 0.1107216;
   Prof_PriceDA.Data[6907] := 0.1107216;
   Prof_PriceDA.Data[6908] := 0.1079028;
   Prof_PriceDA.Data[6909] := 0.1079028;
   Prof_PriceDA.Data[6910] := 0.1079028;
   Prof_PriceDA.Data[6911] := 0.1079028;
   Prof_PriceDA.Data[6912] := 0.1178172;
   Prof_PriceDA.Data[6913] := 0.1178172;
   Prof_PriceDA.Data[6914] := 0.1178172;
   Prof_PriceDA.Data[6915] := 0.1178172;
   Prof_PriceDA.Data[6916] := 0.11448;
   Prof_PriceDA.Data[6917] := 0.11448;
   Prof_PriceDA.Data[6918] := 0.11448;
   Prof_PriceDA.Data[6919] := 0.11448;
   Prof_PriceDA.Data[6920] := 0.114372;
   Prof_PriceDA.Data[6921] := 0.114372;
   Prof_PriceDA.Data[6922] := 0.114372;
   Prof_PriceDA.Data[6923] := 0.114372;
   Prof_PriceDA.Data[6924] := 0.1121364;
   Prof_PriceDA.Data[6925] := 0.1121364;
   Prof_PriceDA.Data[6926] := 0.1121364;
   Prof_PriceDA.Data[6927] := 0.1121364;
   Prof_PriceDA.Data[6928] := 0.113724;
   Prof_PriceDA.Data[6929] := 0.113724;
   Prof_PriceDA.Data[6930] := 0.113724;
   Prof_PriceDA.Data[6931] := 0.113724;
   Prof_PriceDA.Data[6932] := 0.1232928;
   Prof_PriceDA.Data[6933] := 0.1232928;
   Prof_PriceDA.Data[6934] := 0.1232928;
   Prof_PriceDA.Data[6935] := 0.1232928;
   Prof_PriceDA.Data[6936] := 0.1544832;
   Prof_PriceDA.Data[6937] := 0.1544832;
   Prof_PriceDA.Data[6938] := 0.1544832;
   Prof_PriceDA.Data[6939] := 0.1544832;
   Prof_PriceDA.Data[6940] := 0.164646;
   Prof_PriceDA.Data[6941] := 0.164646;
   Prof_PriceDA.Data[6942] := 0.164646;
   Prof_PriceDA.Data[6943] := 0.164646;
   Prof_PriceDA.Data[6944] := 0.1372248;
   Prof_PriceDA.Data[6945] := 0.1372248;
   Prof_PriceDA.Data[6946] := 0.1372248;
   Prof_PriceDA.Data[6947] := 0.1372248;
   Prof_PriceDA.Data[6948] := 0.1197936;
   Prof_PriceDA.Data[6949] := 0.1197936;
   Prof_PriceDA.Data[6950] := 0.1197936;
   Prof_PriceDA.Data[6951] := 0.1197936;
   Prof_PriceDA.Data[6952] := 0.098928;
   Prof_PriceDA.Data[6953] := 0.098928;
   Prof_PriceDA.Data[6954] := 0.098928;
   Prof_PriceDA.Data[6955] := 0.098928;
   Prof_PriceDA.Data[6956] := 0.0945216;
   Prof_PriceDA.Data[6957] := 0.0945216;
   Prof_PriceDA.Data[6958] := 0.0945216;
   Prof_PriceDA.Data[6959] := 0.0945216;
   Prof_PriceDA.Data[6960] := 0.0987228;
   Prof_PriceDA.Data[6961] := 0.0987228;
   Prof_PriceDA.Data[6962] := 0.0987228;
   Prof_PriceDA.Data[6963] := 0.0987228;
   Prof_PriceDA.Data[6964] := 0.098604;
   Prof_PriceDA.Data[6965] := 0.098604;
   Prof_PriceDA.Data[6966] := 0.098604;
   Prof_PriceDA.Data[6967] := 0.098604;
   Prof_PriceDA.Data[6968] := 0.1005372;
   Prof_PriceDA.Data[6969] := 0.1005372;
   Prof_PriceDA.Data[6970] := 0.1005372;
   Prof_PriceDA.Data[6971] := 0.1005372;
   Prof_PriceDA.Data[6972] := 0.1195128;
   Prof_PriceDA.Data[6973] := 0.1195128;
   Prof_PriceDA.Data[6974] := 0.1195128;
   Prof_PriceDA.Data[6975] := 0.1195128;
   Prof_PriceDA.Data[6976] := 0.1374084;
   Prof_PriceDA.Data[6977] := 0.1374084;
   Prof_PriceDA.Data[6978] := 0.1374084;
   Prof_PriceDA.Data[6979] := 0.1374084;
   Prof_PriceDA.Data[6980] := 0.1529388;
   Prof_PriceDA.Data[6981] := 0.1529388;
   Prof_PriceDA.Data[6982] := 0.1529388;
   Prof_PriceDA.Data[6983] := 0.1529388;
   Prof_PriceDA.Data[6984] := 0.1640088;
   Prof_PriceDA.Data[6985] := 0.1640088;
   Prof_PriceDA.Data[6986] := 0.1640088;
   Prof_PriceDA.Data[6987] := 0.1640088;
   Prof_PriceDA.Data[6988] := 0.160002;
   Prof_PriceDA.Data[6989] := 0.160002;
   Prof_PriceDA.Data[6990] := 0.160002;
   Prof_PriceDA.Data[6991] := 0.160002;
   Prof_PriceDA.Data[6992] := 0.1404108;
   Prof_PriceDA.Data[6993] := 0.1404108;
   Prof_PriceDA.Data[6994] := 0.1404108;
   Prof_PriceDA.Data[6995] := 0.1404108;
   Prof_PriceDA.Data[6996] := 0.1203012;
   Prof_PriceDA.Data[6997] := 0.1203012;
   Prof_PriceDA.Data[6998] := 0.1203012;
   Prof_PriceDA.Data[6999] := 0.1203012;
   Prof_PriceDA.Data[7000] := 0.12312;
   Prof_PriceDA.Data[7001] := 0.12312;
   Prof_PriceDA.Data[7002] := 0.12312;
   Prof_PriceDA.Data[7003] := 0.12312;
   Prof_PriceDA.Data[7004] := 0.1135836;
   Prof_PriceDA.Data[7005] := 0.1135836;
   Prof_PriceDA.Data[7006] := 0.1135836;
   Prof_PriceDA.Data[7007] := 0.1135836;
   Prof_PriceDA.Data[7008] := 0.121122;
   Prof_PriceDA.Data[7009] := 0.121122;
   Prof_PriceDA.Data[7010] := 0.121122;
   Prof_PriceDA.Data[7011] := 0.121122;
   Prof_PriceDA.Data[7012] := 0.1113912;
   Prof_PriceDA.Data[7013] := 0.1113912;
   Prof_PriceDA.Data[7014] := 0.1113912;
   Prof_PriceDA.Data[7015] := 0.1113912;
   Prof_PriceDA.Data[7016] := 0.10368;
   Prof_PriceDA.Data[7017] := 0.10368;
   Prof_PriceDA.Data[7018] := 0.10368;
   Prof_PriceDA.Data[7019] := 0.10368;
   Prof_PriceDA.Data[7020] := 0.097092;
   Prof_PriceDA.Data[7021] := 0.097092;
   Prof_PriceDA.Data[7022] := 0.097092;
   Prof_PriceDA.Data[7023] := 0.097092;
   Prof_PriceDA.Data[7024] := 0.093852;
   Prof_PriceDA.Data[7025] := 0.093852;
   Prof_PriceDA.Data[7026] := 0.093852;
   Prof_PriceDA.Data[7027] := 0.093852;
   Prof_PriceDA.Data[7028] := 0.097794;
   Prof_PriceDA.Data[7029] := 0.097794;
   Prof_PriceDA.Data[7030] := 0.097794;
   Prof_PriceDA.Data[7031] := 0.097794;
   Prof_PriceDA.Data[7032] := 0.1047708;
   Prof_PriceDA.Data[7033] := 0.1047708;
   Prof_PriceDA.Data[7034] := 0.1047708;
   Prof_PriceDA.Data[7035] := 0.1047708;
   Prof_PriceDA.Data[7036] := 0.1073736;
   Prof_PriceDA.Data[7037] := 0.1073736;
   Prof_PriceDA.Data[7038] := 0.1073736;
   Prof_PriceDA.Data[7039] := 0.1073736;
   Prof_PriceDA.Data[7040] := 0.0978804;
   Prof_PriceDA.Data[7041] := 0.0978804;
   Prof_PriceDA.Data[7042] := 0.0978804;
   Prof_PriceDA.Data[7043] := 0.0978804;
   Prof_PriceDA.Data[7044] := 0.0824688;
   Prof_PriceDA.Data[7045] := 0.0824688;
   Prof_PriceDA.Data[7046] := 0.0824688;
   Prof_PriceDA.Data[7047] := 0.0824688;
   Prof_PriceDA.Data[7048] := 0.0540432;
   Prof_PriceDA.Data[7049] := 0.0540432;
   Prof_PriceDA.Data[7050] := 0.0540432;
   Prof_PriceDA.Data[7051] := 0.0540432;
   Prof_PriceDA.Data[7052] := 0.016038;
   Prof_PriceDA.Data[7053] := 0.016038;
   Prof_PriceDA.Data[7054] := 0.016038;
   Prof_PriceDA.Data[7055] := 0.016038;
   Prof_PriceDA.Data[7056] := 0.0560736;
   Prof_PriceDA.Data[7057] := 0.0560736;
   Prof_PriceDA.Data[7058] := 0.0560736;
   Prof_PriceDA.Data[7059] := 0.0560736;
   Prof_PriceDA.Data[7060] := 0.05184;
   Prof_PriceDA.Data[7061] := 0.05184;
   Prof_PriceDA.Data[7062] := 0.05184;
   Prof_PriceDA.Data[7063] := 0.05184;
   Prof_PriceDA.Data[7064] := 0.0588708;
   Prof_PriceDA.Data[7065] := 0.0588708;
   Prof_PriceDA.Data[7066] := 0.0588708;
   Prof_PriceDA.Data[7067] := 0.0588708;
   Prof_PriceDA.Data[7068] := 0.0791316;
   Prof_PriceDA.Data[7069] := 0.0791316;
   Prof_PriceDA.Data[7070] := 0.0791316;
   Prof_PriceDA.Data[7071] := 0.0791316;
   Prof_PriceDA.Data[7072] := 0.0940032;
   Prof_PriceDA.Data[7073] := 0.0940032;
   Prof_PriceDA.Data[7074] := 0.0940032;
   Prof_PriceDA.Data[7075] := 0.0940032;
   Prof_PriceDA.Data[7076] := 0.1425492;
   Prof_PriceDA.Data[7077] := 0.1425492;
   Prof_PriceDA.Data[7078] := 0.1425492;
   Prof_PriceDA.Data[7079] := 0.1425492;
   Prof_PriceDA.Data[7080] := 0.15444;
   Prof_PriceDA.Data[7081] := 0.15444;
   Prof_PriceDA.Data[7082] := 0.15444;
   Prof_PriceDA.Data[7083] := 0.15444;
   Prof_PriceDA.Data[7084] := 0.1435968;
   Prof_PriceDA.Data[7085] := 0.1435968;
   Prof_PriceDA.Data[7086] := 0.1435968;
   Prof_PriceDA.Data[7087] := 0.1435968;
   Prof_PriceDA.Data[7088] := 0.1311768;
   Prof_PriceDA.Data[7089] := 0.1311768;
   Prof_PriceDA.Data[7090] := 0.1311768;
   Prof_PriceDA.Data[7091] := 0.1311768;
   Prof_PriceDA.Data[7092] := 0.11718;
   Prof_PriceDA.Data[7093] := 0.11718;
   Prof_PriceDA.Data[7094] := 0.11718;
   Prof_PriceDA.Data[7095] := 0.11718;
   Prof_PriceDA.Data[7096] := 0.1134216;
   Prof_PriceDA.Data[7097] := 0.1134216;
   Prof_PriceDA.Data[7098] := 0.1134216;
   Prof_PriceDA.Data[7099] := 0.1134216;
   Prof_PriceDA.Data[7100] := 0.10287;
   Prof_PriceDA.Data[7101] := 0.10287;
   Prof_PriceDA.Data[7102] := 0.10287;
   Prof_PriceDA.Data[7103] := 0.10287;
   Prof_PriceDA.Data[7104] := 0.0972108;
   Prof_PriceDA.Data[7105] := 0.0972108;
   Prof_PriceDA.Data[7106] := 0.0972108;
   Prof_PriceDA.Data[7107] := 0.0972108;
   Prof_PriceDA.Data[7108] := 0.0926532;
   Prof_PriceDA.Data[7109] := 0.0926532;
   Prof_PriceDA.Data[7110] := 0.0926532;
   Prof_PriceDA.Data[7111] := 0.0926532;
   Prof_PriceDA.Data[7112] := 0.0859896;
   Prof_PriceDA.Data[7113] := 0.0859896;
   Prof_PriceDA.Data[7114] := 0.0859896;
   Prof_PriceDA.Data[7115] := 0.0859896;
   Prof_PriceDA.Data[7116] := 0.0844344;
   Prof_PriceDA.Data[7117] := 0.0844344;
   Prof_PriceDA.Data[7118] := 0.0844344;
   Prof_PriceDA.Data[7119] := 0.0844344;
   Prof_PriceDA.Data[7120] := 0.084888;
   Prof_PriceDA.Data[7121] := 0.084888;
   Prof_PriceDA.Data[7122] := 0.084888;
   Prof_PriceDA.Data[7123] := 0.084888;
   Prof_PriceDA.Data[7124] := 0.0869508;
   Prof_PriceDA.Data[7125] := 0.0869508;
   Prof_PriceDA.Data[7126] := 0.0869508;
   Prof_PriceDA.Data[7127] := 0.0869508;
   Prof_PriceDA.Data[7128] := 0.0919512;
   Prof_PriceDA.Data[7129] := 0.0919512;
   Prof_PriceDA.Data[7130] := 0.0919512;
   Prof_PriceDA.Data[7131] := 0.0919512;
   Prof_PriceDA.Data[7132] := 0.0886356;
   Prof_PriceDA.Data[7133] := 0.0886356;
   Prof_PriceDA.Data[7134] := 0.0886356;
   Prof_PriceDA.Data[7135] := 0.0886356;
   Prof_PriceDA.Data[7136] := 0.084186;
   Prof_PriceDA.Data[7137] := 0.084186;
   Prof_PriceDA.Data[7138] := 0.084186;
   Prof_PriceDA.Data[7139] := 0.084186;
   Prof_PriceDA.Data[7140] := 0.0742608;
   Prof_PriceDA.Data[7141] := 0.0742608;
   Prof_PriceDA.Data[7142] := 0.0742608;
   Prof_PriceDA.Data[7143] := 0.0742608;
   Prof_PriceDA.Data[7144] := 0.0340956;
   Prof_PriceDA.Data[7145] := 0.0340956;
   Prof_PriceDA.Data[7146] := 0.0340956;
   Prof_PriceDA.Data[7147] := 0.0340956;
   Prof_PriceDA.Data[7148] := 0.0137268;
   Prof_PriceDA.Data[7149] := 0.0137268;
   Prof_PriceDA.Data[7150] := 0.0137268;
   Prof_PriceDA.Data[7151] := 0.0137268;
   Prof_PriceDA.Data[7152] := 0.0090072;
   Prof_PriceDA.Data[7153] := 0.0090072;
   Prof_PriceDA.Data[7154] := 0.0090072;
   Prof_PriceDA.Data[7155] := 0.0090072;
   Prof_PriceDA.Data[7156] := 0.0057564;
   Prof_PriceDA.Data[7157] := 0.0057564;
   Prof_PriceDA.Data[7158] := 0.0057564;
   Prof_PriceDA.Data[7159] := 0.0057564;
   Prof_PriceDA.Data[7160] := 0.0104112;
   Prof_PriceDA.Data[7161] := 0.0104112;
   Prof_PriceDA.Data[7162] := 0.0104112;
   Prof_PriceDA.Data[7163] := 0.0104112;
   Prof_PriceDA.Data[7164] := 0.03348;
   Prof_PriceDA.Data[7165] := 0.03348;
   Prof_PriceDA.Data[7166] := 0.03348;
   Prof_PriceDA.Data[7167] := 0.03348;
   Prof_PriceDA.Data[7168] := 0.0786024;
   Prof_PriceDA.Data[7169] := 0.0786024;
   Prof_PriceDA.Data[7170] := 0.0786024;
   Prof_PriceDA.Data[7171] := 0.0786024;
   Prof_PriceDA.Data[7172] := 0.1285416;
   Prof_PriceDA.Data[7173] := 0.1285416;
   Prof_PriceDA.Data[7174] := 0.1285416;
   Prof_PriceDA.Data[7175] := 0.1285416;
   Prof_PriceDA.Data[7176] := 0.1432188;
   Prof_PriceDA.Data[7177] := 0.1432188;
   Prof_PriceDA.Data[7178] := 0.1432188;
   Prof_PriceDA.Data[7179] := 0.1432188;
   Prof_PriceDA.Data[7180] := 0.1512;
   Prof_PriceDA.Data[7181] := 0.1512;
   Prof_PriceDA.Data[7182] := 0.1512;
   Prof_PriceDA.Data[7183] := 0.1512;
   Prof_PriceDA.Data[7184] := 0.1364364;
   Prof_PriceDA.Data[7185] := 0.1364364;
   Prof_PriceDA.Data[7186] := 0.1364364;
   Prof_PriceDA.Data[7187] := 0.1364364;
   Prof_PriceDA.Data[7188] := 0.1175796;
   Prof_PriceDA.Data[7189] := 0.1175796;
   Prof_PriceDA.Data[7190] := 0.1175796;
   Prof_PriceDA.Data[7191] := 0.1175796;
   Prof_PriceDA.Data[7192] := 0.1102248;
   Prof_PriceDA.Data[7193] := 0.1102248;
   Prof_PriceDA.Data[7194] := 0.1102248;
   Prof_PriceDA.Data[7195] := 0.1102248;
   Prof_PriceDA.Data[7196] := 0.088614;
   Prof_PriceDA.Data[7197] := 0.088614;
   Prof_PriceDA.Data[7198] := 0.088614;
   Prof_PriceDA.Data[7199] := 0.088614;
   Prof_PriceDA.Data[7200] := 0.0892296;
   Prof_PriceDA.Data[7201] := 0.0892296;
   Prof_PriceDA.Data[7202] := 0.0892296;
   Prof_PriceDA.Data[7203] := 0.0892296;
   Prof_PriceDA.Data[7204] := 0.0895212;
   Prof_PriceDA.Data[7205] := 0.0895212;
   Prof_PriceDA.Data[7206] := 0.0895212;
   Prof_PriceDA.Data[7207] := 0.0895212;
   Prof_PriceDA.Data[7208] := 0.0872208;
   Prof_PriceDA.Data[7209] := 0.0872208;
   Prof_PriceDA.Data[7210] := 0.0872208;
   Prof_PriceDA.Data[7211] := 0.0872208;
   Prof_PriceDA.Data[7212] := 0.0873828;
   Prof_PriceDA.Data[7213] := 0.0873828;
   Prof_PriceDA.Data[7214] := 0.0873828;
   Prof_PriceDA.Data[7215] := 0.0873828;
   Prof_PriceDA.Data[7216] := 0.092718;
   Prof_PriceDA.Data[7217] := 0.092718;
   Prof_PriceDA.Data[7218] := 0.092718;
   Prof_PriceDA.Data[7219] := 0.092718;
   Prof_PriceDA.Data[7220] := 0.111564;
   Prof_PriceDA.Data[7221] := 0.111564;
   Prof_PriceDA.Data[7222] := 0.111564;
   Prof_PriceDA.Data[7223] := 0.111564;
   Prof_PriceDA.Data[7224] := 0.1459944;
   Prof_PriceDA.Data[7225] := 0.1459944;
   Prof_PriceDA.Data[7226] := 0.1459944;
   Prof_PriceDA.Data[7227] := 0.1459944;
   Prof_PriceDA.Data[7228] := 0.1650996;
   Prof_PriceDA.Data[7229] := 0.1650996;
   Prof_PriceDA.Data[7230] := 0.1650996;
   Prof_PriceDA.Data[7231] := 0.1650996;
   Prof_PriceDA.Data[7232] := 0.1475496;
   Prof_PriceDA.Data[7233] := 0.1475496;
   Prof_PriceDA.Data[7234] := 0.1475496;
   Prof_PriceDA.Data[7235] := 0.1475496;
   Prof_PriceDA.Data[7236] := 0.1150524;
   Prof_PriceDA.Data[7237] := 0.1150524;
   Prof_PriceDA.Data[7238] := 0.1150524;
   Prof_PriceDA.Data[7239] := 0.1150524;
   Prof_PriceDA.Data[7240] := 0.0911736;
   Prof_PriceDA.Data[7241] := 0.0911736;
   Prof_PriceDA.Data[7242] := 0.0911736;
   Prof_PriceDA.Data[7243] := 0.0911736;
   Prof_PriceDA.Data[7244] := 0.0838188;
   Prof_PriceDA.Data[7245] := 0.0838188;
   Prof_PriceDA.Data[7246] := 0.0838188;
   Prof_PriceDA.Data[7247] := 0.0838188;
   Prof_PriceDA.Data[7248] := 0.0725976;
   Prof_PriceDA.Data[7249] := 0.0725976;
   Prof_PriceDA.Data[7250] := 0.0725976;
   Prof_PriceDA.Data[7251] := 0.0725976;
   Prof_PriceDA.Data[7252] := 0.0486756;
   Prof_PriceDA.Data[7253] := 0.0486756;
   Prof_PriceDA.Data[7254] := 0.0486756;
   Prof_PriceDA.Data[7255] := 0.0486756;
   Prof_PriceDA.Data[7256] := 0.0543132;
   Prof_PriceDA.Data[7257] := 0.0543132;
   Prof_PriceDA.Data[7258] := 0.0543132;
   Prof_PriceDA.Data[7259] := 0.0543132;
   Prof_PriceDA.Data[7260] := 0.0770472;
   Prof_PriceDA.Data[7261] := 0.0770472;
   Prof_PriceDA.Data[7262] := 0.0770472;
   Prof_PriceDA.Data[7263] := 0.0770472;
   Prof_PriceDA.Data[7264] := 0.1122876;
   Prof_PriceDA.Data[7265] := 0.1122876;
   Prof_PriceDA.Data[7266] := 0.1122876;
   Prof_PriceDA.Data[7267] := 0.1122876;
   Prof_PriceDA.Data[7268] := 0.1642572;
   Prof_PriceDA.Data[7269] := 0.1642572;
   Prof_PriceDA.Data[7270] := 0.1642572;
   Prof_PriceDA.Data[7271] := 0.1642572;
   Prof_PriceDA.Data[7272] := 0.1824984;
   Prof_PriceDA.Data[7273] := 0.1824984;
   Prof_PriceDA.Data[7274] := 0.1824984;
   Prof_PriceDA.Data[7275] := 0.1824984;
   Prof_PriceDA.Data[7276] := 0.1836;
   Prof_PriceDA.Data[7277] := 0.1836;
   Prof_PriceDA.Data[7278] := 0.1836;
   Prof_PriceDA.Data[7279] := 0.1836;
   Prof_PriceDA.Data[7280] := 0.15282;
   Prof_PriceDA.Data[7281] := 0.15282;
   Prof_PriceDA.Data[7282] := 0.15282;
   Prof_PriceDA.Data[7283] := 0.15282;
   Prof_PriceDA.Data[7284] := 0.1292544;
   Prof_PriceDA.Data[7285] := 0.1292544;
   Prof_PriceDA.Data[7286] := 0.1292544;
   Prof_PriceDA.Data[7287] := 0.1292544;
   Prof_PriceDA.Data[7288] := 0.1171152;
   Prof_PriceDA.Data[7289] := 0.1171152;
   Prof_PriceDA.Data[7290] := 0.1171152;
   Prof_PriceDA.Data[7291] := 0.1171152;
   Prof_PriceDA.Data[7292] := 0.10098;
   Prof_PriceDA.Data[7293] := 0.10098;
   Prof_PriceDA.Data[7294] := 0.10098;
   Prof_PriceDA.Data[7295] := 0.10098;
   Prof_PriceDA.Data[7296] := 0.099576;
   Prof_PriceDA.Data[7297] := 0.099576;
   Prof_PriceDA.Data[7298] := 0.099576;
   Prof_PriceDA.Data[7299] := 0.099576;
   Prof_PriceDA.Data[7300] := 0.0971892;
   Prof_PriceDA.Data[7301] := 0.0971892;
   Prof_PriceDA.Data[7302] := 0.0971892;
   Prof_PriceDA.Data[7303] := 0.0971892;
   Prof_PriceDA.Data[7304] := 0.1000404;
   Prof_PriceDA.Data[7305] := 0.1000404;
   Prof_PriceDA.Data[7306] := 0.1000404;
   Prof_PriceDA.Data[7307] := 0.1000404;
   Prof_PriceDA.Data[7308] := 0.096876;
   Prof_PriceDA.Data[7309] := 0.096876;
   Prof_PriceDA.Data[7310] := 0.096876;
   Prof_PriceDA.Data[7311] := 0.096876;
   Prof_PriceDA.Data[7312] := 0.103248;
   Prof_PriceDA.Data[7313] := 0.103248;
   Prof_PriceDA.Data[7314] := 0.103248;
   Prof_PriceDA.Data[7315] := 0.103248;
   Prof_PriceDA.Data[7316] := 0.1221804;
   Prof_PriceDA.Data[7317] := 0.1221804;
   Prof_PriceDA.Data[7318] := 0.1221804;
   Prof_PriceDA.Data[7319] := 0.1221804;
   Prof_PriceDA.Data[7320] := 0.1527228;
   Prof_PriceDA.Data[7321] := 0.1527228;
   Prof_PriceDA.Data[7322] := 0.1527228;
   Prof_PriceDA.Data[7323] := 0.1527228;
   Prof_PriceDA.Data[7324] := 0.1476144;
   Prof_PriceDA.Data[7325] := 0.1476144;
   Prof_PriceDA.Data[7326] := 0.1476144;
   Prof_PriceDA.Data[7327] := 0.1476144;
   Prof_PriceDA.Data[7328] := 0.0788184;
   Prof_PriceDA.Data[7329] := 0.0788184;
   Prof_PriceDA.Data[7330] := 0.0788184;
   Prof_PriceDA.Data[7331] := 0.0788184;
   Prof_PriceDA.Data[7332] := 0.0556524;
   Prof_PriceDA.Data[7333] := 0.0556524;
   Prof_PriceDA.Data[7334] := 0.0556524;
   Prof_PriceDA.Data[7335] := 0.0556524;
   Prof_PriceDA.Data[7336] := 0.033966;
   Prof_PriceDA.Data[7337] := 0.033966;
   Prof_PriceDA.Data[7338] := 0.033966;
   Prof_PriceDA.Data[7339] := 0.033966;
   Prof_PriceDA.Data[7340] := 0.0033156;
   Prof_PriceDA.Data[7341] := 0.0033156;
   Prof_PriceDA.Data[7342] := 0.0033156;
   Prof_PriceDA.Data[7343] := 0.0033156;
   Prof_PriceDA.Data[7344] := 0.0044496;
   Prof_PriceDA.Data[7345] := 0.0044496;
   Prof_PriceDA.Data[7346] := 0.0044496;
   Prof_PriceDA.Data[7347] := 0.0044496;
   Prof_PriceDA.Data[7348] := 0.0034992;
   Prof_PriceDA.Data[7349] := 0.0034992;
   Prof_PriceDA.Data[7350] := 0.0034992;
   Prof_PriceDA.Data[7351] := 0.0034992;
   Prof_PriceDA.Data[7352] := 0.0080676;
   Prof_PriceDA.Data[7353] := 0.0080676;
   Prof_PriceDA.Data[7354] := 0.0080676;
   Prof_PriceDA.Data[7355] := 0.0080676;
   Prof_PriceDA.Data[7356] := 0.0745524;
   Prof_PriceDA.Data[7357] := 0.0745524;
   Prof_PriceDA.Data[7358] := 0.0745524;
   Prof_PriceDA.Data[7359] := 0.0745524;
   Prof_PriceDA.Data[7360] := 0.1153116;
   Prof_PriceDA.Data[7361] := 0.1153116;
   Prof_PriceDA.Data[7362] := 0.1153116;
   Prof_PriceDA.Data[7363] := 0.1153116;
   Prof_PriceDA.Data[7364] := 0.1616328;
   Prof_PriceDA.Data[7365] := 0.1616328;
   Prof_PriceDA.Data[7366] := 0.1616328;
   Prof_PriceDA.Data[7367] := 0.1616328;
   Prof_PriceDA.Data[7368] := 0.18495;
   Prof_PriceDA.Data[7369] := 0.18495;
   Prof_PriceDA.Data[7370] := 0.18495;
   Prof_PriceDA.Data[7371] := 0.18495;
   Prof_PriceDA.Data[7372] := 0.178416;
   Prof_PriceDA.Data[7373] := 0.178416;
   Prof_PriceDA.Data[7374] := 0.178416;
   Prof_PriceDA.Data[7375] := 0.178416;
   Prof_PriceDA.Data[7376] := 0.1556388;
   Prof_PriceDA.Data[7377] := 0.1556388;
   Prof_PriceDA.Data[7378] := 0.1556388;
   Prof_PriceDA.Data[7379] := 0.1556388;
   Prof_PriceDA.Data[7380] := 0.1349568;
   Prof_PriceDA.Data[7381] := 0.1349568;
   Prof_PriceDA.Data[7382] := 0.1349568;
   Prof_PriceDA.Data[7383] := 0.1349568;
   Prof_PriceDA.Data[7384] := 0.1285092;
   Prof_PriceDA.Data[7385] := 0.1285092;
   Prof_PriceDA.Data[7386] := 0.1285092;
   Prof_PriceDA.Data[7387] := 0.1285092;
   Prof_PriceDA.Data[7388] := 0.1130112;
   Prof_PriceDA.Data[7389] := 0.1130112;
   Prof_PriceDA.Data[7390] := 0.1130112;
   Prof_PriceDA.Data[7391] := 0.1130112;
   Prof_PriceDA.Data[7392] := 0.1197396;
   Prof_PriceDA.Data[7393] := 0.1197396;
   Prof_PriceDA.Data[7394] := 0.1197396;
   Prof_PriceDA.Data[7395] := 0.1197396;
   Prof_PriceDA.Data[7396] := 0.1151928;
   Prof_PriceDA.Data[7397] := 0.1151928;
   Prof_PriceDA.Data[7398] := 0.1151928;
   Prof_PriceDA.Data[7399] := 0.1151928;
   Prof_PriceDA.Data[7400] := 0.113292;
   Prof_PriceDA.Data[7401] := 0.113292;
   Prof_PriceDA.Data[7402] := 0.113292;
   Prof_PriceDA.Data[7403] := 0.113292;
   Prof_PriceDA.Data[7404] := 0.1126548;
   Prof_PriceDA.Data[7405] := 0.1126548;
   Prof_PriceDA.Data[7406] := 0.1126548;
   Prof_PriceDA.Data[7407] := 0.1126548;
   Prof_PriceDA.Data[7408] := 0.1180764;
   Prof_PriceDA.Data[7409] := 0.1180764;
   Prof_PriceDA.Data[7410] := 0.1180764;
   Prof_PriceDA.Data[7411] := 0.1180764;
   Prof_PriceDA.Data[7412] := 0.138024;
   Prof_PriceDA.Data[7413] := 0.138024;
   Prof_PriceDA.Data[7414] := 0.138024;
   Prof_PriceDA.Data[7415] := 0.138024;
   Prof_PriceDA.Data[7416] := 0.1770012;
   Prof_PriceDA.Data[7417] := 0.1770012;
   Prof_PriceDA.Data[7418] := 0.1770012;
   Prof_PriceDA.Data[7419] := 0.1770012;
   Prof_PriceDA.Data[7420] := 0.1575828;
   Prof_PriceDA.Data[7421] := 0.1575828;
   Prof_PriceDA.Data[7422] := 0.1575828;
   Prof_PriceDA.Data[7423] := 0.1575828;
   Prof_PriceDA.Data[7424] := 0.1099116;
   Prof_PriceDA.Data[7425] := 0.1099116;
   Prof_PriceDA.Data[7426] := 0.1099116;
   Prof_PriceDA.Data[7427] := 0.1099116;
   Prof_PriceDA.Data[7428] := 0.0314172;
   Prof_PriceDA.Data[7429] := 0.0314172;
   Prof_PriceDA.Data[7430] := 0.0314172;
   Prof_PriceDA.Data[7431] := 0.0314172;
   Prof_PriceDA.Data[7432] := 0.0230472;
   Prof_PriceDA.Data[7433] := 0.0230472;
   Prof_PriceDA.Data[7434] := 0.0230472;
   Prof_PriceDA.Data[7435] := 0.0230472;
   Prof_PriceDA.Data[7436] := 0.0017064;
   Prof_PriceDA.Data[7437] := 0.0017064;
   Prof_PriceDA.Data[7438] := 0.0017064;
   Prof_PriceDA.Data[7439] := 0.0017064;
   Prof_PriceDA.Data[7440] := 0.0002052;
   Prof_PriceDA.Data[7441] := 0.0002052;
   Prof_PriceDA.Data[7442] := 0.0002052;
   Prof_PriceDA.Data[7443] := 0.0002052;
   Prof_PriceDA.Data[7444] := 0.001404;
   Prof_PriceDA.Data[7445] := 0.001404;
   Prof_PriceDA.Data[7446] := 0.001404;
   Prof_PriceDA.Data[7447] := 0.001404;
   Prof_PriceDA.Data[7448] := 0.0042444;
   Prof_PriceDA.Data[7449] := 0.0042444;
   Prof_PriceDA.Data[7450] := 0.0042444;
   Prof_PriceDA.Data[7451] := 0.0042444;
   Prof_PriceDA.Data[7452] := 0.07425;
   Prof_PriceDA.Data[7453] := 0.07425;
   Prof_PriceDA.Data[7454] := 0.07425;
   Prof_PriceDA.Data[7455] := 0.07425;
   Prof_PriceDA.Data[7456] := 0.1289088;
   Prof_PriceDA.Data[7457] := 0.1289088;
   Prof_PriceDA.Data[7458] := 0.1289088;
   Prof_PriceDA.Data[7459] := 0.1289088;
   Prof_PriceDA.Data[7460] := 0.1772928;
   Prof_PriceDA.Data[7461] := 0.1772928;
   Prof_PriceDA.Data[7462] := 0.1772928;
   Prof_PriceDA.Data[7463] := 0.1772928;
   Prof_PriceDA.Data[7464] := 0.2667708;
   Prof_PriceDA.Data[7465] := 0.2667708;
   Prof_PriceDA.Data[7466] := 0.2667708;
   Prof_PriceDA.Data[7467] := 0.2667708;
   Prof_PriceDA.Data[7468] := 0.2296512;
   Prof_PriceDA.Data[7469] := 0.2296512;
   Prof_PriceDA.Data[7470] := 0.2296512;
   Prof_PriceDA.Data[7471] := 0.2296512;
   Prof_PriceDA.Data[7472] := 0.1785348;
   Prof_PriceDA.Data[7473] := 0.1785348;
   Prof_PriceDA.Data[7474] := 0.1785348;
   Prof_PriceDA.Data[7475] := 0.1785348;
   Prof_PriceDA.Data[7476] := 0.1571184;
   Prof_PriceDA.Data[7477] := 0.1571184;
   Prof_PriceDA.Data[7478] := 0.1571184;
   Prof_PriceDA.Data[7479] := 0.1571184;
   Prof_PriceDA.Data[7480] := 0.1424952;
   Prof_PriceDA.Data[7481] := 0.1424952;
   Prof_PriceDA.Data[7482] := 0.1424952;
   Prof_PriceDA.Data[7483] := 0.1424952;
   Prof_PriceDA.Data[7484] := 0.1250316;
   Prof_PriceDA.Data[7485] := 0.1250316;
   Prof_PriceDA.Data[7486] := 0.1250316;
   Prof_PriceDA.Data[7487] := 0.1250316;
   Prof_PriceDA.Data[7488] := 0.1358532;
   Prof_PriceDA.Data[7489] := 0.1358532;
   Prof_PriceDA.Data[7490] := 0.1358532;
   Prof_PriceDA.Data[7491] := 0.1358532;
   Prof_PriceDA.Data[7492] := 0.119772;
   Prof_PriceDA.Data[7493] := 0.119772;
   Prof_PriceDA.Data[7494] := 0.119772;
   Prof_PriceDA.Data[7495] := 0.119772;
   Prof_PriceDA.Data[7496] := 0.1138968;
   Prof_PriceDA.Data[7497] := 0.1138968;
   Prof_PriceDA.Data[7498] := 0.1138968;
   Prof_PriceDA.Data[7499] := 0.1138968;
   Prof_PriceDA.Data[7500] := 0.1154304;
   Prof_PriceDA.Data[7501] := 0.1154304;
   Prof_PriceDA.Data[7502] := 0.1154304;
   Prof_PriceDA.Data[7503] := 0.1154304;
   Prof_PriceDA.Data[7504] := 0.1230444;
   Prof_PriceDA.Data[7505] := 0.1230444;
   Prof_PriceDA.Data[7506] := 0.1230444;
   Prof_PriceDA.Data[7507] := 0.1230444;
   Prof_PriceDA.Data[7508] := 0.141642;
   Prof_PriceDA.Data[7509] := 0.141642;
   Prof_PriceDA.Data[7510] := 0.141642;
   Prof_PriceDA.Data[7511] := 0.141642;
   Prof_PriceDA.Data[7512] := 0.1664928;
   Prof_PriceDA.Data[7513] := 0.1664928;
   Prof_PriceDA.Data[7514] := 0.1664928;
   Prof_PriceDA.Data[7515] := 0.1664928;
   Prof_PriceDA.Data[7516] := 0.1559628;
   Prof_PriceDA.Data[7517] := 0.1559628;
   Prof_PriceDA.Data[7518] := 0.1559628;
   Prof_PriceDA.Data[7519] := 0.1559628;
   Prof_PriceDA.Data[7520] := 0.1072116;
   Prof_PriceDA.Data[7521] := 0.1072116;
   Prof_PriceDA.Data[7522] := 0.1072116;
   Prof_PriceDA.Data[7523] := 0.1072116;
   Prof_PriceDA.Data[7524] := 0.087264;
   Prof_PriceDA.Data[7525] := 0.087264;
   Prof_PriceDA.Data[7526] := 0.087264;
   Prof_PriceDA.Data[7527] := 0.087264;
   Prof_PriceDA.Data[7528] := 0.0393336;
   Prof_PriceDA.Data[7529] := 0.0393336;
   Prof_PriceDA.Data[7530] := 0.0393336;
   Prof_PriceDA.Data[7531] := 0.0393336;
   Prof_PriceDA.Data[7532] := 0.0036936;
   Prof_PriceDA.Data[7533] := 0.0036936;
   Prof_PriceDA.Data[7534] := 0.0036936;
   Prof_PriceDA.Data[7535] := 0.0036936;
   Prof_PriceDA.Data[7536] := 0.0004644;
   Prof_PriceDA.Data[7537] := 0.0004644;
   Prof_PriceDA.Data[7538] := 0.0004644;
   Prof_PriceDA.Data[7539] := 0.0004644;
   Prof_PriceDA.Data[7540] := 0.000702;
   Prof_PriceDA.Data[7541] := 0.000702;
   Prof_PriceDA.Data[7542] := 0.000702;
   Prof_PriceDA.Data[7543] := 0.000702;
   Prof_PriceDA.Data[7544] := 0.0190728;
   Prof_PriceDA.Data[7545] := 0.0190728;
   Prof_PriceDA.Data[7546] := 0.0190728;
   Prof_PriceDA.Data[7547] := 0.0190728;
   Prof_PriceDA.Data[7548] := 0.0910548;
   Prof_PriceDA.Data[7549] := 0.0910548;
   Prof_PriceDA.Data[7550] := 0.0910548;
   Prof_PriceDA.Data[7551] := 0.0910548;
   Prof_PriceDA.Data[7552] := 0.1377324;
   Prof_PriceDA.Data[7553] := 0.1377324;
   Prof_PriceDA.Data[7554] := 0.1377324;
   Prof_PriceDA.Data[7555] := 0.1377324;
   Prof_PriceDA.Data[7556] := 0.1914516;
   Prof_PriceDA.Data[7557] := 0.1914516;
   Prof_PriceDA.Data[7558] := 0.1914516;
   Prof_PriceDA.Data[7559] := 0.1914516;
   Prof_PriceDA.Data[7560] := 0.2737044;
   Prof_PriceDA.Data[7561] := 0.2737044;
   Prof_PriceDA.Data[7562] := 0.2737044;
   Prof_PriceDA.Data[7563] := 0.2737044;
   Prof_PriceDA.Data[7564] := 0.2508084;
   Prof_PriceDA.Data[7565] := 0.2508084;
   Prof_PriceDA.Data[7566] := 0.2508084;
   Prof_PriceDA.Data[7567] := 0.2508084;
   Prof_PriceDA.Data[7568] := 0.1867536;
   Prof_PriceDA.Data[7569] := 0.1867536;
   Prof_PriceDA.Data[7570] := 0.1867536;
   Prof_PriceDA.Data[7571] := 0.1867536;
   Prof_PriceDA.Data[7572] := 0.1605096;
   Prof_PriceDA.Data[7573] := 0.1605096;
   Prof_PriceDA.Data[7574] := 0.1605096;
   Prof_PriceDA.Data[7575] := 0.1605096;
   Prof_PriceDA.Data[7576] := 0.1471608;
   Prof_PriceDA.Data[7577] := 0.1471608;
   Prof_PriceDA.Data[7578] := 0.1471608;
   Prof_PriceDA.Data[7579] := 0.1471608;
   Prof_PriceDA.Data[7580] := 0.137484;
   Prof_PriceDA.Data[7581] := 0.137484;
   Prof_PriceDA.Data[7582] := 0.137484;
   Prof_PriceDA.Data[7583] := 0.137484;
   Prof_PriceDA.Data[7584] := 0.1430244;
   Prof_PriceDA.Data[7585] := 0.1430244;
   Prof_PriceDA.Data[7586] := 0.1430244;
   Prof_PriceDA.Data[7587] := 0.1430244;
   Prof_PriceDA.Data[7588] := 0.132408;
   Prof_PriceDA.Data[7589] := 0.132408;
   Prof_PriceDA.Data[7590] := 0.132408;
   Prof_PriceDA.Data[7591] := 0.132408;
   Prof_PriceDA.Data[7592] := 0.1289088;
   Prof_PriceDA.Data[7593] := 0.1289088;
   Prof_PriceDA.Data[7594] := 0.1289088;
   Prof_PriceDA.Data[7595] := 0.1289088;
   Prof_PriceDA.Data[7596] := 0.1239192;
   Prof_PriceDA.Data[7597] := 0.1239192;
   Prof_PriceDA.Data[7598] := 0.1239192;
   Prof_PriceDA.Data[7599] := 0.1239192;
   Prof_PriceDA.Data[7600] := 0.128898;
   Prof_PriceDA.Data[7601] := 0.128898;
   Prof_PriceDA.Data[7602] := 0.128898;
   Prof_PriceDA.Data[7603] := 0.128898;
   Prof_PriceDA.Data[7604] := 0.1521288;
   Prof_PriceDA.Data[7605] := 0.1521288;
   Prof_PriceDA.Data[7606] := 0.1521288;
   Prof_PriceDA.Data[7607] := 0.1521288;
   Prof_PriceDA.Data[7608] := 0.1841832;
   Prof_PriceDA.Data[7609] := 0.1841832;
   Prof_PriceDA.Data[7610] := 0.1841832;
   Prof_PriceDA.Data[7611] := 0.1841832;
   Prof_PriceDA.Data[7612] := 0.1653588;
   Prof_PriceDA.Data[7613] := 0.1653588;
   Prof_PriceDA.Data[7614] := 0.1653588;
   Prof_PriceDA.Data[7615] := 0.1653588;
   Prof_PriceDA.Data[7616] := 0.1232388;
   Prof_PriceDA.Data[7617] := 0.1232388;
   Prof_PriceDA.Data[7618] := 0.1232388;
   Prof_PriceDA.Data[7619] := 0.1232388;
   Prof_PriceDA.Data[7620] := 0.0808056;
   Prof_PriceDA.Data[7621] := 0.0808056;
   Prof_PriceDA.Data[7622] := 0.0808056;
   Prof_PriceDA.Data[7623] := 0.0808056;
   Prof_PriceDA.Data[7624] := 0.0430488;
   Prof_PriceDA.Data[7625] := 0.0430488;
   Prof_PriceDA.Data[7626] := 0.0430488;
   Prof_PriceDA.Data[7627] := 0.0430488;
   Prof_PriceDA.Data[7628] := 0.0079056;
   Prof_PriceDA.Data[7629] := 0.0079056;
   Prof_PriceDA.Data[7630] := 0.0079056;
   Prof_PriceDA.Data[7631] := 0.0079056;
   Prof_PriceDA.Data[7632] := 0.00189;
   Prof_PriceDA.Data[7633] := 0.00189;
   Prof_PriceDA.Data[7634] := 0.00189;
   Prof_PriceDA.Data[7635] := 0.00189;
   Prof_PriceDA.Data[7636] := 0.0002376;
   Prof_PriceDA.Data[7637] := 0.0002376;
   Prof_PriceDA.Data[7638] := 0.0002376;
   Prof_PriceDA.Data[7639] := 0.0002376;
   Prof_PriceDA.Data[7640] := 0.0067608;
   Prof_PriceDA.Data[7641] := 0.0067608;
   Prof_PriceDA.Data[7642] := 0.0067608;
   Prof_PriceDA.Data[7643] := 0.0067608;
   Prof_PriceDA.Data[7644] := 0.0624348;
   Prof_PriceDA.Data[7645] := 0.0624348;
   Prof_PriceDA.Data[7646] := 0.0624348;
   Prof_PriceDA.Data[7647] := 0.0624348;
   Prof_PriceDA.Data[7648] := 0.1274616;
   Prof_PriceDA.Data[7649] := 0.1274616;
   Prof_PriceDA.Data[7650] := 0.1274616;
   Prof_PriceDA.Data[7651] := 0.1274616;
   Prof_PriceDA.Data[7652] := 0.1607364;
   Prof_PriceDA.Data[7653] := 0.1607364;
   Prof_PriceDA.Data[7654] := 0.1607364;
   Prof_PriceDA.Data[7655] := 0.1607364;
   Prof_PriceDA.Data[7656] := 0.2246508;
   Prof_PriceDA.Data[7657] := 0.2246508;
   Prof_PriceDA.Data[7658] := 0.2246508;
   Prof_PriceDA.Data[7659] := 0.2246508;
   Prof_PriceDA.Data[7660] := 0.1900584;
   Prof_PriceDA.Data[7661] := 0.1900584;
   Prof_PriceDA.Data[7662] := 0.1900584;
   Prof_PriceDA.Data[7663] := 0.1900584;
   Prof_PriceDA.Data[7664] := 0.1624212;
   Prof_PriceDA.Data[7665] := 0.1624212;
   Prof_PriceDA.Data[7666] := 0.1624212;
   Prof_PriceDA.Data[7667] := 0.1624212;
   Prof_PriceDA.Data[7668] := 0.1486404;
   Prof_PriceDA.Data[7669] := 0.1486404;
   Prof_PriceDA.Data[7670] := 0.1486404;
   Prof_PriceDA.Data[7671] := 0.1486404;
   Prof_PriceDA.Data[7672] := 0.132354;
   Prof_PriceDA.Data[7673] := 0.132354;
   Prof_PriceDA.Data[7674] := 0.132354;
   Prof_PriceDA.Data[7675] := 0.132354;
   Prof_PriceDA.Data[7676] := 0.1172556;
   Prof_PriceDA.Data[7677] := 0.1172556;
   Prof_PriceDA.Data[7678] := 0.1172556;
   Prof_PriceDA.Data[7679] := 0.1172556;
   Prof_PriceDA.Data[7680] := 0.106812;
   Prof_PriceDA.Data[7681] := 0.106812;
   Prof_PriceDA.Data[7682] := 0.106812;
   Prof_PriceDA.Data[7683] := 0.106812;
   Prof_PriceDA.Data[7684] := 0.0965088;
   Prof_PriceDA.Data[7685] := 0.0965088;
   Prof_PriceDA.Data[7686] := 0.0965088;
   Prof_PriceDA.Data[7687] := 0.0965088;
   Prof_PriceDA.Data[7688] := 0.1034424;
   Prof_PriceDA.Data[7689] := 0.1034424;
   Prof_PriceDA.Data[7690] := 0.1034424;
   Prof_PriceDA.Data[7691] := 0.1034424;
   Prof_PriceDA.Data[7692] := 0.1046304;
   Prof_PriceDA.Data[7693] := 0.1046304;
   Prof_PriceDA.Data[7694] := 0.1046304;
   Prof_PriceDA.Data[7695] := 0.1046304;
   Prof_PriceDA.Data[7696] := 0.1058292;
   Prof_PriceDA.Data[7697] := 0.1058292;
   Prof_PriceDA.Data[7698] := 0.1058292;
   Prof_PriceDA.Data[7699] := 0.1058292;
   Prof_PriceDA.Data[7700] := 0.1103976;
   Prof_PriceDA.Data[7701] := 0.1103976;
   Prof_PriceDA.Data[7702] := 0.1103976;
   Prof_PriceDA.Data[7703] := 0.1103976;
   Prof_PriceDA.Data[7704] := 0.0961416;
   Prof_PriceDA.Data[7705] := 0.0961416;
   Prof_PriceDA.Data[7706] := 0.0961416;
   Prof_PriceDA.Data[7707] := 0.0961416;
   Prof_PriceDA.Data[7708] := 0.076086;
   Prof_PriceDA.Data[7709] := 0.076086;
   Prof_PriceDA.Data[7710] := 0.076086;
   Prof_PriceDA.Data[7711] := 0.076086;
   Prof_PriceDA.Data[7712] := 0.0631044;
   Prof_PriceDA.Data[7713] := 0.0631044;
   Prof_PriceDA.Data[7714] := 0.0631044;
   Prof_PriceDA.Data[7715] := 0.0631044;
   Prof_PriceDA.Data[7716] := 0.0527472;
   Prof_PriceDA.Data[7717] := 0.0527472;
   Prof_PriceDA.Data[7718] := 0.0527472;
   Prof_PriceDA.Data[7719] := 0.0527472;
   Prof_PriceDA.Data[7720] := 0.023598;
   Prof_PriceDA.Data[7721] := 0.023598;
   Prof_PriceDA.Data[7722] := 0.023598;
   Prof_PriceDA.Data[7723] := 0.023598;
   Prof_PriceDA.Data[7724] := 0.0159948;
   Prof_PriceDA.Data[7725] := 0.0159948;
   Prof_PriceDA.Data[7726] := 0.0159948;
   Prof_PriceDA.Data[7727] := 0.0159948;
   Prof_PriceDA.Data[7728] := 0.046926;
   Prof_PriceDA.Data[7729] := 0.046926;
   Prof_PriceDA.Data[7730] := 0.046926;
   Prof_PriceDA.Data[7731] := 0.046926;
   Prof_PriceDA.Data[7732] := 0.0540972;
   Prof_PriceDA.Data[7733] := 0.0540972;
   Prof_PriceDA.Data[7734] := 0.0540972;
   Prof_PriceDA.Data[7735] := 0.0540972;
   Prof_PriceDA.Data[7736] := 0.0613224;
   Prof_PriceDA.Data[7737] := 0.0613224;
   Prof_PriceDA.Data[7738] := 0.0613224;
   Prof_PriceDA.Data[7739] := 0.0613224;
   Prof_PriceDA.Data[7740] := 0.0924372;
   Prof_PriceDA.Data[7741] := 0.0924372;
   Prof_PriceDA.Data[7742] := 0.0924372;
   Prof_PriceDA.Data[7743] := 0.0924372;
   Prof_PriceDA.Data[7744] := 0.1254852;
   Prof_PriceDA.Data[7745] := 0.1254852;
   Prof_PriceDA.Data[7746] := 0.1254852;
   Prof_PriceDA.Data[7747] := 0.1254852;
   Prof_PriceDA.Data[7748] := 0.1314252;
   Prof_PriceDA.Data[7749] := 0.1314252;
   Prof_PriceDA.Data[7750] := 0.1314252;
   Prof_PriceDA.Data[7751] := 0.1314252;
   Prof_PriceDA.Data[7752] := 0.1388988;
   Prof_PriceDA.Data[7753] := 0.1388988;
   Prof_PriceDA.Data[7754] := 0.1388988;
   Prof_PriceDA.Data[7755] := 0.1388988;
   Prof_PriceDA.Data[7756] := 0.1359504;
   Prof_PriceDA.Data[7757] := 0.1359504;
   Prof_PriceDA.Data[7758] := 0.1359504;
   Prof_PriceDA.Data[7759] := 0.1359504;
   Prof_PriceDA.Data[7760] := 0.1250316;
   Prof_PriceDA.Data[7761] := 0.1250316;
   Prof_PriceDA.Data[7762] := 0.1250316;
   Prof_PriceDA.Data[7763] := 0.1250316;
   Prof_PriceDA.Data[7764] := 0.0847152;
   Prof_PriceDA.Data[7765] := 0.0847152;
   Prof_PriceDA.Data[7766] := 0.0847152;
   Prof_PriceDA.Data[7767] := 0.0847152;
   Prof_PriceDA.Data[7768] := 0.081108;
   Prof_PriceDA.Data[7769] := 0.081108;
   Prof_PriceDA.Data[7770] := 0.081108;
   Prof_PriceDA.Data[7771] := 0.081108;
   Prof_PriceDA.Data[7772] := 0.06696;
   Prof_PriceDA.Data[7773] := 0.06696;
   Prof_PriceDA.Data[7774] := 0.06696;
   Prof_PriceDA.Data[7775] := 0.06696;
   Prof_PriceDA.Data[7776] := 0.0401004;
   Prof_PriceDA.Data[7777] := 0.0401004;
   Prof_PriceDA.Data[7778] := 0.0401004;
   Prof_PriceDA.Data[7779] := 0.0401004;
   Prof_PriceDA.Data[7780] := 0.03915;
   Prof_PriceDA.Data[7781] := 0.03915;
   Prof_PriceDA.Data[7782] := 0.03915;
   Prof_PriceDA.Data[7783] := 0.03915;
   Prof_PriceDA.Data[7784] := 0.0478116;
   Prof_PriceDA.Data[7785] := 0.0478116;
   Prof_PriceDA.Data[7786] := 0.0478116;
   Prof_PriceDA.Data[7787] := 0.0478116;
   Prof_PriceDA.Data[7788] := 0.0467424;
   Prof_PriceDA.Data[7789] := 0.0467424;
   Prof_PriceDA.Data[7790] := 0.0467424;
   Prof_PriceDA.Data[7791] := 0.0467424;
   Prof_PriceDA.Data[7792] := 0.0470232;
   Prof_PriceDA.Data[7793] := 0.0470232;
   Prof_PriceDA.Data[7794] := 0.0470232;
   Prof_PriceDA.Data[7795] := 0.0470232;
   Prof_PriceDA.Data[7796] := 0.0467316;
   Prof_PriceDA.Data[7797] := 0.0467316;
   Prof_PriceDA.Data[7798] := 0.0467316;
   Prof_PriceDA.Data[7799] := 0.0467316;
   Prof_PriceDA.Data[7800] := 0.0483192;
   Prof_PriceDA.Data[7801] := 0.0483192;
   Prof_PriceDA.Data[7802] := 0.0483192;
   Prof_PriceDA.Data[7803] := 0.0483192;
   Prof_PriceDA.Data[7804] := 0.041256;
   Prof_PriceDA.Data[7805] := 0.041256;
   Prof_PriceDA.Data[7806] := 0.041256;
   Prof_PriceDA.Data[7807] := 0.041256;
   Prof_PriceDA.Data[7808] := 0.0276156;
   Prof_PriceDA.Data[7809] := 0.0276156;
   Prof_PriceDA.Data[7810] := 0.0276156;
   Prof_PriceDA.Data[7811] := 0.0276156;
   Prof_PriceDA.Data[7812] := 0.0231984;
   Prof_PriceDA.Data[7813] := 0.0231984;
   Prof_PriceDA.Data[7814] := 0.0231984;
   Prof_PriceDA.Data[7815] := 0.0231984;
   Prof_PriceDA.Data[7816] := 0.0148824;
   Prof_PriceDA.Data[7817] := 0.0148824;
   Prof_PriceDA.Data[7818] := 0.0148824;
   Prof_PriceDA.Data[7819] := 0.0148824;
   Prof_PriceDA.Data[7820] := 0.010368;
   Prof_PriceDA.Data[7821] := 0.010368;
   Prof_PriceDA.Data[7822] := 0.010368;
   Prof_PriceDA.Data[7823] := 0.010368;
   Prof_PriceDA.Data[7824] := 0.0145692;
   Prof_PriceDA.Data[7825] := 0.0145692;
   Prof_PriceDA.Data[7826] := 0.0145692;
   Prof_PriceDA.Data[7827] := 0.0145692;
   Prof_PriceDA.Data[7828] := 0.0054108;
   Prof_PriceDA.Data[7829] := 0.0054108;
   Prof_PriceDA.Data[7830] := 0.0054108;
   Prof_PriceDA.Data[7831] := 0.0054108;
   Prof_PriceDA.Data[7832] := 0.0123768;
   Prof_PriceDA.Data[7833] := 0.0123768;
   Prof_PriceDA.Data[7834] := 0.0123768;
   Prof_PriceDA.Data[7835] := 0.0123768;
   Prof_PriceDA.Data[7836] := 0.0467208;
   Prof_PriceDA.Data[7837] := 0.0467208;
   Prof_PriceDA.Data[7838] := 0.0467208;
   Prof_PriceDA.Data[7839] := 0.0467208;
   Prof_PriceDA.Data[7840] := 0.097092;
   Prof_PriceDA.Data[7841] := 0.097092;
   Prof_PriceDA.Data[7842] := 0.097092;
   Prof_PriceDA.Data[7843] := 0.097092;
   Prof_PriceDA.Data[7844] := 0.1409076;
   Prof_PriceDA.Data[7845] := 0.1409076;
   Prof_PriceDA.Data[7846] := 0.1409076;
   Prof_PriceDA.Data[7847] := 0.1409076;
   Prof_PriceDA.Data[7848] := 0.1566756;
   Prof_PriceDA.Data[7849] := 0.1566756;
   Prof_PriceDA.Data[7850] := 0.1566756;
   Prof_PriceDA.Data[7851] := 0.1566756;
   Prof_PriceDA.Data[7852] := 0.1554228;
   Prof_PriceDA.Data[7853] := 0.1554228;
   Prof_PriceDA.Data[7854] := 0.1554228;
   Prof_PriceDA.Data[7855] := 0.1554228;
   Prof_PriceDA.Data[7856] := 0.151632;
   Prof_PriceDA.Data[7857] := 0.151632;
   Prof_PriceDA.Data[7858] := 0.151632;
   Prof_PriceDA.Data[7859] := 0.151632;
   Prof_PriceDA.Data[7860] := 0.1417932;
   Prof_PriceDA.Data[7861] := 0.1417932;
   Prof_PriceDA.Data[7862] := 0.1417932;
   Prof_PriceDA.Data[7863] := 0.1417932;
   Prof_PriceDA.Data[7864] := 0.1374084;
   Prof_PriceDA.Data[7865] := 0.1374084;
   Prof_PriceDA.Data[7866] := 0.1374084;
   Prof_PriceDA.Data[7867] := 0.1374084;
   Prof_PriceDA.Data[7868] := 0.1233792;
   Prof_PriceDA.Data[7869] := 0.1233792;
   Prof_PriceDA.Data[7870] := 0.1233792;
   Prof_PriceDA.Data[7871] := 0.1233792;
   Prof_PriceDA.Data[7872] := 0.1183032;
   Prof_PriceDA.Data[7873] := 0.1183032;
   Prof_PriceDA.Data[7874] := 0.1183032;
   Prof_PriceDA.Data[7875] := 0.1183032;
   Prof_PriceDA.Data[7876] := 0.11637;
   Prof_PriceDA.Data[7877] := 0.11637;
   Prof_PriceDA.Data[7878] := 0.11637;
   Prof_PriceDA.Data[7879] := 0.11637;
   Prof_PriceDA.Data[7880] := 0.1103112;
   Prof_PriceDA.Data[7881] := 0.1103112;
   Prof_PriceDA.Data[7882] := 0.1103112;
   Prof_PriceDA.Data[7883] := 0.1103112;
   Prof_PriceDA.Data[7884] := 0.107298;
   Prof_PriceDA.Data[7885] := 0.107298;
   Prof_PriceDA.Data[7886] := 0.107298;
   Prof_PriceDA.Data[7887] := 0.107298;
   Prof_PriceDA.Data[7888] := 0.1109052;
   Prof_PriceDA.Data[7889] := 0.1109052;
   Prof_PriceDA.Data[7890] := 0.1109052;
   Prof_PriceDA.Data[7891] := 0.1109052;
   Prof_PriceDA.Data[7892] := 0.1302696;
   Prof_PriceDA.Data[7893] := 0.1302696;
   Prof_PriceDA.Data[7894] := 0.1302696;
   Prof_PriceDA.Data[7895] := 0.1302696;
   Prof_PriceDA.Data[7896] := 0.1545156;
   Prof_PriceDA.Data[7897] := 0.1545156;
   Prof_PriceDA.Data[7898] := 0.1545156;
   Prof_PriceDA.Data[7899] := 0.1545156;
   Prof_PriceDA.Data[7900] := 0.1774008;
   Prof_PriceDA.Data[7901] := 0.1774008;
   Prof_PriceDA.Data[7902] := 0.1774008;
   Prof_PriceDA.Data[7903] := 0.1774008;
   Prof_PriceDA.Data[7904] := 0.1754136;
   Prof_PriceDA.Data[7905] := 0.1754136;
   Prof_PriceDA.Data[7906] := 0.1754136;
   Prof_PriceDA.Data[7907] := 0.1754136;
   Prof_PriceDA.Data[7908] := 0.1472364;
   Prof_PriceDA.Data[7909] := 0.1472364;
   Prof_PriceDA.Data[7910] := 0.1472364;
   Prof_PriceDA.Data[7911] := 0.1472364;
   Prof_PriceDA.Data[7912] := 0.1205388;
   Prof_PriceDA.Data[7913] := 0.1205388;
   Prof_PriceDA.Data[7914] := 0.1205388;
   Prof_PriceDA.Data[7915] := 0.1205388;
   Prof_PriceDA.Data[7916] := 0.1193184;
   Prof_PriceDA.Data[7917] := 0.1193184;
   Prof_PriceDA.Data[7918] := 0.1193184;
   Prof_PriceDA.Data[7919] := 0.1193184;
   Prof_PriceDA.Data[7920] := 0.113616;
   Prof_PriceDA.Data[7921] := 0.113616;
   Prof_PriceDA.Data[7922] := 0.113616;
   Prof_PriceDA.Data[7923] := 0.113616;
   Prof_PriceDA.Data[7924] := 0.1166832;
   Prof_PriceDA.Data[7925] := 0.1166832;
   Prof_PriceDA.Data[7926] := 0.1166832;
   Prof_PriceDA.Data[7927] := 0.1166832;
   Prof_PriceDA.Data[7928] := 0.1260144;
   Prof_PriceDA.Data[7929] := 0.1260144;
   Prof_PriceDA.Data[7930] := 0.1260144;
   Prof_PriceDA.Data[7931] := 0.1260144;
   Prof_PriceDA.Data[7932] := 0.1354752;
   Prof_PriceDA.Data[7933] := 0.1354752;
   Prof_PriceDA.Data[7934] := 0.1354752;
   Prof_PriceDA.Data[7935] := 0.1354752;
   Prof_PriceDA.Data[7936] := 0.1469664;
   Prof_PriceDA.Data[7937] := 0.1469664;
   Prof_PriceDA.Data[7938] := 0.1469664;
   Prof_PriceDA.Data[7939] := 0.1469664;
   Prof_PriceDA.Data[7940] := 0.1676052;
   Prof_PriceDA.Data[7941] := 0.1676052;
   Prof_PriceDA.Data[7942] := 0.1676052;
   Prof_PriceDA.Data[7943] := 0.1676052;
   Prof_PriceDA.Data[7944] := 0.225018;
   Prof_PriceDA.Data[7945] := 0.225018;
   Prof_PriceDA.Data[7946] := 0.225018;
   Prof_PriceDA.Data[7947] := 0.225018;
   Prof_PriceDA.Data[7948] := 0.2084832;
   Prof_PriceDA.Data[7949] := 0.2084832;
   Prof_PriceDA.Data[7950] := 0.2084832;
   Prof_PriceDA.Data[7951] := 0.2084832;
   Prof_PriceDA.Data[7952] := 0.1749708;
   Prof_PriceDA.Data[7953] := 0.1749708;
   Prof_PriceDA.Data[7954] := 0.1749708;
   Prof_PriceDA.Data[7955] := 0.1749708;
   Prof_PriceDA.Data[7956] := 0.150984;
   Prof_PriceDA.Data[7957] := 0.150984;
   Prof_PriceDA.Data[7958] := 0.150984;
   Prof_PriceDA.Data[7959] := 0.150984;
   Prof_PriceDA.Data[7960] := 0.1370196;
   Prof_PriceDA.Data[7961] := 0.1370196;
   Prof_PriceDA.Data[7962] := 0.1370196;
   Prof_PriceDA.Data[7963] := 0.1370196;
   Prof_PriceDA.Data[7964] := 0.1251072;
   Prof_PriceDA.Data[7965] := 0.1251072;
   Prof_PriceDA.Data[7966] := 0.1251072;
   Prof_PriceDA.Data[7967] := 0.1251072;
   Prof_PriceDA.Data[7968] := 0.10989;
   Prof_PriceDA.Data[7969] := 0.10989;
   Prof_PriceDA.Data[7970] := 0.10989;
   Prof_PriceDA.Data[7971] := 0.10989;
   Prof_PriceDA.Data[7972] := 0.1109808;
   Prof_PriceDA.Data[7973] := 0.1109808;
   Prof_PriceDA.Data[7974] := 0.1109808;
   Prof_PriceDA.Data[7975] := 0.1109808;
   Prof_PriceDA.Data[7976] := 0.1094148;
   Prof_PriceDA.Data[7977] := 0.1094148;
   Prof_PriceDA.Data[7978] := 0.1094148;
   Prof_PriceDA.Data[7979] := 0.1094148;
   Prof_PriceDA.Data[7980] := 0.1137564;
   Prof_PriceDA.Data[7981] := 0.1137564;
   Prof_PriceDA.Data[7982] := 0.1137564;
   Prof_PriceDA.Data[7983] := 0.1137564;
   Prof_PriceDA.Data[7984] := 0.113076;
   Prof_PriceDA.Data[7985] := 0.113076;
   Prof_PriceDA.Data[7986] := 0.113076;
   Prof_PriceDA.Data[7987] := 0.113076;
   Prof_PriceDA.Data[7988] := 0.1185732;
   Prof_PriceDA.Data[7989] := 0.1185732;
   Prof_PriceDA.Data[7990] := 0.1185732;
   Prof_PriceDA.Data[7991] := 0.1185732;
   Prof_PriceDA.Data[7992] := 0.1511568;
   Prof_PriceDA.Data[7993] := 0.1511568;
   Prof_PriceDA.Data[7994] := 0.1511568;
   Prof_PriceDA.Data[7995] := 0.1511568;
   Prof_PriceDA.Data[7996] := 0.1553904;
   Prof_PriceDA.Data[7997] := 0.1553904;
   Prof_PriceDA.Data[7998] := 0.1553904;
   Prof_PriceDA.Data[7999] := 0.1553904;
   Prof_PriceDA.Data[8000] := 0.1502604;
   Prof_PriceDA.Data[8001] := 0.1502604;
   Prof_PriceDA.Data[8002] := 0.1502604;
   Prof_PriceDA.Data[8003] := 0.1502604;
   Prof_PriceDA.Data[8004] := 0.12474;
   Prof_PriceDA.Data[8005] := 0.12474;
   Prof_PriceDA.Data[8006] := 0.12474;
   Prof_PriceDA.Data[8007] := 0.12474;
   Prof_PriceDA.Data[8008] := 0.11718;
   Prof_PriceDA.Data[8009] := 0.11718;
   Prof_PriceDA.Data[8010] := 0.11718;
   Prof_PriceDA.Data[8011] := 0.11718;
   Prof_PriceDA.Data[8012] := 0.1110024;
   Prof_PriceDA.Data[8013] := 0.1110024;
   Prof_PriceDA.Data[8014] := 0.1110024;
   Prof_PriceDA.Data[8015] := 0.1110024;
   Prof_PriceDA.Data[8016] := 0.1050516;
   Prof_PriceDA.Data[8017] := 0.1050516;
   Prof_PriceDA.Data[8018] := 0.1050516;
   Prof_PriceDA.Data[8019] := 0.1050516;
   Prof_PriceDA.Data[8020] := 0.1064772;
   Prof_PriceDA.Data[8021] := 0.1064772;
   Prof_PriceDA.Data[8022] := 0.1064772;
   Prof_PriceDA.Data[8023] := 0.1064772;
   Prof_PriceDA.Data[8024] := 0.1191672;
   Prof_PriceDA.Data[8025] := 0.1191672;
   Prof_PriceDA.Data[8026] := 0.1191672;
   Prof_PriceDA.Data[8027] := 0.1191672;
   Prof_PriceDA.Data[8028] := 0.1322028;
   Prof_PriceDA.Data[8029] := 0.1322028;
   Prof_PriceDA.Data[8030] := 0.1322028;
   Prof_PriceDA.Data[8031] := 0.1322028;
   Prof_PriceDA.Data[8032] := 0.1511568;
   Prof_PriceDA.Data[8033] := 0.1511568;
   Prof_PriceDA.Data[8034] := 0.1511568;
   Prof_PriceDA.Data[8035] := 0.1511568;
   Prof_PriceDA.Data[8036] := 0.15525;
   Prof_PriceDA.Data[8037] := 0.15525;
   Prof_PriceDA.Data[8038] := 0.15525;
   Prof_PriceDA.Data[8039] := 0.15525;
   Prof_PriceDA.Data[8040] := 0.1925208;
   Prof_PriceDA.Data[8041] := 0.1925208;
   Prof_PriceDA.Data[8042] := 0.1925208;
   Prof_PriceDA.Data[8043] := 0.1925208;
   Prof_PriceDA.Data[8044] := 0.1871856;
   Prof_PriceDA.Data[8045] := 0.1871856;
   Prof_PriceDA.Data[8046] := 0.1871856;
   Prof_PriceDA.Data[8047] := 0.1871856;
   Prof_PriceDA.Data[8048] := 0.160488;
   Prof_PriceDA.Data[8049] := 0.160488;
   Prof_PriceDA.Data[8050] := 0.160488;
   Prof_PriceDA.Data[8051] := 0.160488;
   Prof_PriceDA.Data[8052] := 0.1487268;
   Prof_PriceDA.Data[8053] := 0.1487268;
   Prof_PriceDA.Data[8054] := 0.1487268;
   Prof_PriceDA.Data[8055] := 0.1487268;
   Prof_PriceDA.Data[8056] := 0.1365984;
   Prof_PriceDA.Data[8057] := 0.1365984;
   Prof_PriceDA.Data[8058] := 0.1365984;
   Prof_PriceDA.Data[8059] := 0.1365984;
   Prof_PriceDA.Data[8060] := 0.110214;
   Prof_PriceDA.Data[8061] := 0.110214;
   Prof_PriceDA.Data[8062] := 0.110214;
   Prof_PriceDA.Data[8063] := 0.110214;
   Prof_PriceDA.Data[8064] := 0.1091016;
   Prof_PriceDA.Data[8065] := 0.1091016;
   Prof_PriceDA.Data[8066] := 0.1091016;
   Prof_PriceDA.Data[8067] := 0.1091016;
   Prof_PriceDA.Data[8068] := 0.106596;
   Prof_PriceDA.Data[8069] := 0.106596;
   Prof_PriceDA.Data[8070] := 0.106596;
   Prof_PriceDA.Data[8071] := 0.106596;
   Prof_PriceDA.Data[8072] := 0.1064016;
   Prof_PriceDA.Data[8073] := 0.1064016;
   Prof_PriceDA.Data[8074] := 0.1064016;
   Prof_PriceDA.Data[8075] := 0.1064016;
   Prof_PriceDA.Data[8076] := 0.1079244;
   Prof_PriceDA.Data[8077] := 0.1079244;
   Prof_PriceDA.Data[8078] := 0.1079244;
   Prof_PriceDA.Data[8079] := 0.1079244;
   Prof_PriceDA.Data[8080] := 0.1107216;
   Prof_PriceDA.Data[8081] := 0.1107216;
   Prof_PriceDA.Data[8082] := 0.1107216;
   Prof_PriceDA.Data[8083] := 0.1107216;
   Prof_PriceDA.Data[8084] := 0.1205388;
   Prof_PriceDA.Data[8085] := 0.1205388;
   Prof_PriceDA.Data[8086] := 0.1205388;
   Prof_PriceDA.Data[8087] := 0.1205388;
   Prof_PriceDA.Data[8088] := 0.1464264;
   Prof_PriceDA.Data[8089] := 0.1464264;
   Prof_PriceDA.Data[8090] := 0.1464264;
   Prof_PriceDA.Data[8091] := 0.1464264;
   Prof_PriceDA.Data[8092] := 0.1543536;
   Prof_PriceDA.Data[8093] := 0.1543536;
   Prof_PriceDA.Data[8094] := 0.1543536;
   Prof_PriceDA.Data[8095] := 0.1543536;
   Prof_PriceDA.Data[8096] := 0.1490616;
   Prof_PriceDA.Data[8097] := 0.1490616;
   Prof_PriceDA.Data[8098] := 0.1490616;
   Prof_PriceDA.Data[8099] := 0.1490616;
   Prof_PriceDA.Data[8100] := 0.1211652;
   Prof_PriceDA.Data[8101] := 0.1211652;
   Prof_PriceDA.Data[8102] := 0.1211652;
   Prof_PriceDA.Data[8103] := 0.1211652;
   Prof_PriceDA.Data[8104] := 0.1083348;
   Prof_PriceDA.Data[8105] := 0.1083348;
   Prof_PriceDA.Data[8106] := 0.1083348;
   Prof_PriceDA.Data[8107] := 0.1083348;
   Prof_PriceDA.Data[8108] := 0.1047708;
   Prof_PriceDA.Data[8109] := 0.1047708;
   Prof_PriceDA.Data[8110] := 0.1047708;
   Prof_PriceDA.Data[8111] := 0.1047708;
   Prof_PriceDA.Data[8112] := 0.1027296;
   Prof_PriceDA.Data[8113] := 0.1027296;
   Prof_PriceDA.Data[8114] := 0.1027296;
   Prof_PriceDA.Data[8115] := 0.1027296;
   Prof_PriceDA.Data[8116] := 0.091908;
   Prof_PriceDA.Data[8117] := 0.091908;
   Prof_PriceDA.Data[8118] := 0.091908;
   Prof_PriceDA.Data[8119] := 0.091908;
   Prof_PriceDA.Data[8120] := 0.1026864;
   Prof_PriceDA.Data[8121] := 0.1026864;
   Prof_PriceDA.Data[8122] := 0.1026864;
   Prof_PriceDA.Data[8123] := 0.1026864;
   Prof_PriceDA.Data[8124] := 0.110538;
   Prof_PriceDA.Data[8125] := 0.110538;
   Prof_PriceDA.Data[8126] := 0.110538;
   Prof_PriceDA.Data[8127] := 0.110538;
   Prof_PriceDA.Data[8128] := 0.127116;
   Prof_PriceDA.Data[8129] := 0.127116;
   Prof_PriceDA.Data[8130] := 0.127116;
   Prof_PriceDA.Data[8131] := 0.127116;
   Prof_PriceDA.Data[8132] := 0.154818;
   Prof_PriceDA.Data[8133] := 0.154818;
   Prof_PriceDA.Data[8134] := 0.154818;
   Prof_PriceDA.Data[8135] := 0.154818;
   Prof_PriceDA.Data[8136] := 0.1812996;
   Prof_PriceDA.Data[8137] := 0.1812996;
   Prof_PriceDA.Data[8138] := 0.1812996;
   Prof_PriceDA.Data[8139] := 0.1812996;
   Prof_PriceDA.Data[8140] := 0.1863648;
   Prof_PriceDA.Data[8141] := 0.1863648;
   Prof_PriceDA.Data[8142] := 0.1863648;
   Prof_PriceDA.Data[8143] := 0.1863648;
   Prof_PriceDA.Data[8144] := 0.1700028;
   Prof_PriceDA.Data[8145] := 0.1700028;
   Prof_PriceDA.Data[8146] := 0.1700028;
   Prof_PriceDA.Data[8147] := 0.1700028;
   Prof_PriceDA.Data[8148] := 0.142668;
   Prof_PriceDA.Data[8149] := 0.142668;
   Prof_PriceDA.Data[8150] := 0.142668;
   Prof_PriceDA.Data[8151] := 0.142668;
   Prof_PriceDA.Data[8152] := 0.1342008;
   Prof_PriceDA.Data[8153] := 0.1342008;
   Prof_PriceDA.Data[8154] := 0.1342008;
   Prof_PriceDA.Data[8155] := 0.1342008;
   Prof_PriceDA.Data[8156] := 0.1196856;
   Prof_PriceDA.Data[8157] := 0.1196856;
   Prof_PriceDA.Data[8158] := 0.1196856;
   Prof_PriceDA.Data[8159] := 0.1196856;
   Prof_PriceDA.Data[8160] := 0.1138104;
   Prof_PriceDA.Data[8161] := 0.1138104;
   Prof_PriceDA.Data[8162] := 0.1138104;
   Prof_PriceDA.Data[8163] := 0.1138104;
   Prof_PriceDA.Data[8164] := 0.1077084;
   Prof_PriceDA.Data[8165] := 0.1077084;
   Prof_PriceDA.Data[8166] := 0.1077084;
   Prof_PriceDA.Data[8167] := 0.1077084;
   Prof_PriceDA.Data[8168] := 0.1057968;
   Prof_PriceDA.Data[8169] := 0.1057968;
   Prof_PriceDA.Data[8170] := 0.1057968;
   Prof_PriceDA.Data[8171] := 0.1057968;
   Prof_PriceDA.Data[8172] := 0.1071468;
   Prof_PriceDA.Data[8173] := 0.1071468;
   Prof_PriceDA.Data[8174] := 0.1071468;
   Prof_PriceDA.Data[8175] := 0.1071468;
   Prof_PriceDA.Data[8176] := 0.1059372;
   Prof_PriceDA.Data[8177] := 0.1059372;
   Prof_PriceDA.Data[8178] := 0.1059372;
   Prof_PriceDA.Data[8179] := 0.1059372;
   Prof_PriceDA.Data[8180] := 0.1139292;
   Prof_PriceDA.Data[8181] := 0.1139292;
   Prof_PriceDA.Data[8182] := 0.1139292;
   Prof_PriceDA.Data[8183] := 0.1139292;
   Prof_PriceDA.Data[8184] := 0.1418364;
   Prof_PriceDA.Data[8185] := 0.1418364;
   Prof_PriceDA.Data[8186] := 0.1418364;
   Prof_PriceDA.Data[8187] := 0.1418364;
   Prof_PriceDA.Data[8188] := 0.15228;
   Prof_PriceDA.Data[8189] := 0.15228;
   Prof_PriceDA.Data[8190] := 0.15228;
   Prof_PriceDA.Data[8191] := 0.15228;
   Prof_PriceDA.Data[8192] := 0.13338;
   Prof_PriceDA.Data[8193] := 0.13338;
   Prof_PriceDA.Data[8194] := 0.13338;
   Prof_PriceDA.Data[8195] := 0.13338;
   Prof_PriceDA.Data[8196] := 0.0971136;
   Prof_PriceDA.Data[8197] := 0.0971136;
   Prof_PriceDA.Data[8198] := 0.0971136;
   Prof_PriceDA.Data[8199] := 0.0971136;
   Prof_PriceDA.Data[8200] := 0.0874692;
   Prof_PriceDA.Data[8201] := 0.0874692;
   Prof_PriceDA.Data[8202] := 0.0874692;
   Prof_PriceDA.Data[8203] := 0.0874692;
   Prof_PriceDA.Data[8204] := 0.0493992;
   Prof_PriceDA.Data[8205] := 0.0493992;
   Prof_PriceDA.Data[8206] := 0.0493992;
   Prof_PriceDA.Data[8207] := 0.0493992;
   Prof_PriceDA.Data[8208] := 0.04212;
   Prof_PriceDA.Data[8209] := 0.04212;
   Prof_PriceDA.Data[8210] := 0.04212;
   Prof_PriceDA.Data[8211] := 0.04212;
   Prof_PriceDA.Data[8212] := 0.0297;
   Prof_PriceDA.Data[8213] := 0.0297;
   Prof_PriceDA.Data[8214] := 0.0297;
   Prof_PriceDA.Data[8215] := 0.0297;
   Prof_PriceDA.Data[8216] := 0.0637956;
   Prof_PriceDA.Data[8217] := 0.0637956;
   Prof_PriceDA.Data[8218] := 0.0637956;
   Prof_PriceDA.Data[8219] := 0.0637956;
   Prof_PriceDA.Data[8220] := 0.0911844;
   Prof_PriceDA.Data[8221] := 0.0911844;
   Prof_PriceDA.Data[8222] := 0.0911844;
   Prof_PriceDA.Data[8223] := 0.0911844;
   Prof_PriceDA.Data[8224] := 0.1082484;
   Prof_PriceDA.Data[8225] := 0.1082484;
   Prof_PriceDA.Data[8226] := 0.1082484;
   Prof_PriceDA.Data[8227] := 0.1082484;
   Prof_PriceDA.Data[8228] := 0.1454544;
   Prof_PriceDA.Data[8229] := 0.1454544;
   Prof_PriceDA.Data[8230] := 0.1454544;
   Prof_PriceDA.Data[8231] := 0.1454544;
   Prof_PriceDA.Data[8232] := 0.1713312;
   Prof_PriceDA.Data[8233] := 0.1713312;
   Prof_PriceDA.Data[8234] := 0.1713312;
   Prof_PriceDA.Data[8235] := 0.1713312;
   Prof_PriceDA.Data[8236] := 0.1830816;
   Prof_PriceDA.Data[8237] := 0.1830816;
   Prof_PriceDA.Data[8238] := 0.1830816;
   Prof_PriceDA.Data[8239] := 0.1830816;
   Prof_PriceDA.Data[8240] := 0.1533384;
   Prof_PriceDA.Data[8241] := 0.1533384;
   Prof_PriceDA.Data[8242] := 0.1533384;
   Prof_PriceDA.Data[8243] := 0.1533384;
   Prof_PriceDA.Data[8244] := 0.1351404;
   Prof_PriceDA.Data[8245] := 0.1351404;
   Prof_PriceDA.Data[8246] := 0.1351404;
   Prof_PriceDA.Data[8247] := 0.1351404;
   Prof_PriceDA.Data[8248] := 0.12285;
   Prof_PriceDA.Data[8249] := 0.12285;
   Prof_PriceDA.Data[8250] := 0.12285;
   Prof_PriceDA.Data[8251] := 0.12285;
   Prof_PriceDA.Data[8252] := 0.109512;
   Prof_PriceDA.Data[8253] := 0.109512;
   Prof_PriceDA.Data[8254] := 0.109512;
   Prof_PriceDA.Data[8255] := 0.109512;
   Prof_PriceDA.Data[8256] := 0.099144;
   Prof_PriceDA.Data[8257] := 0.099144;
   Prof_PriceDA.Data[8258] := 0.099144;
   Prof_PriceDA.Data[8259] := 0.099144;
   Prof_PriceDA.Data[8260] := 0.08586;
   Prof_PriceDA.Data[8261] := 0.08586;
   Prof_PriceDA.Data[8262] := 0.08586;
   Prof_PriceDA.Data[8263] := 0.08586;
   Prof_PriceDA.Data[8264] := 0.0853416;
   Prof_PriceDA.Data[8265] := 0.0853416;
   Prof_PriceDA.Data[8266] := 0.0853416;
   Prof_PriceDA.Data[8267] := 0.0853416;
   Prof_PriceDA.Data[8268] := 0.0862488;
   Prof_PriceDA.Data[8269] := 0.0862488;
   Prof_PriceDA.Data[8270] := 0.0862488;
   Prof_PriceDA.Data[8271] := 0.0862488;
   Prof_PriceDA.Data[8272] := 0.086778;
   Prof_PriceDA.Data[8273] := 0.086778;
   Prof_PriceDA.Data[8274] := 0.086778;
   Prof_PriceDA.Data[8275] := 0.086778;
   Prof_PriceDA.Data[8276] := 0.1185948;
   Prof_PriceDA.Data[8277] := 0.1185948;
   Prof_PriceDA.Data[8278] := 0.1185948;
   Prof_PriceDA.Data[8279] := 0.1185948;
   Prof_PriceDA.Data[8280] := 0.141156;
   Prof_PriceDA.Data[8281] := 0.141156;
   Prof_PriceDA.Data[8282] := 0.141156;
   Prof_PriceDA.Data[8283] := 0.141156;
   Prof_PriceDA.Data[8284] := 0.131976;
   Prof_PriceDA.Data[8285] := 0.131976;
   Prof_PriceDA.Data[8286] := 0.131976;
   Prof_PriceDA.Data[8287] := 0.131976;
   Prof_PriceDA.Data[8288] := 0.1102464;
   Prof_PriceDA.Data[8289] := 0.1102464;
   Prof_PriceDA.Data[8290] := 0.1102464;
   Prof_PriceDA.Data[8291] := 0.1102464;
   Prof_PriceDA.Data[8292] := 0.0834624;
   Prof_PriceDA.Data[8293] := 0.0834624;
   Prof_PriceDA.Data[8294] := 0.0834624;
   Prof_PriceDA.Data[8295] := 0.0834624;
   Prof_PriceDA.Data[8296] := 0.073872;
   Prof_PriceDA.Data[8297] := 0.073872;
   Prof_PriceDA.Data[8298] := 0.073872;
   Prof_PriceDA.Data[8299] := 0.073872;
   Prof_PriceDA.Data[8300] := 0.0550908;
   Prof_PriceDA.Data[8301] := 0.0550908;
   Prof_PriceDA.Data[8302] := 0.0550908;
   Prof_PriceDA.Data[8303] := 0.0550908;
   Prof_PriceDA.Data[8304] := 0.0735588;
   Prof_PriceDA.Data[8305] := 0.0735588;
   Prof_PriceDA.Data[8306] := 0.0735588;
   Prof_PriceDA.Data[8307] := 0.0735588;
   Prof_PriceDA.Data[8308] := 0.081054;
   Prof_PriceDA.Data[8309] := 0.081054;
   Prof_PriceDA.Data[8310] := 0.081054;
   Prof_PriceDA.Data[8311] := 0.081054;
   Prof_PriceDA.Data[8312] := 0.0810432;
   Prof_PriceDA.Data[8313] := 0.0810432;
   Prof_PriceDA.Data[8314] := 0.0810432;
   Prof_PriceDA.Data[8315] := 0.0810432;
   Prof_PriceDA.Data[8316] := 0.112914;
   Prof_PriceDA.Data[8317] := 0.112914;
   Prof_PriceDA.Data[8318] := 0.112914;
   Prof_PriceDA.Data[8319] := 0.112914;
   Prof_PriceDA.Data[8320] := 0.1191132;
   Prof_PriceDA.Data[8321] := 0.1191132;
   Prof_PriceDA.Data[8322] := 0.1191132;
   Prof_PriceDA.Data[8323] := 0.1191132;
   Prof_PriceDA.Data[8324] := 0.1475928;
   Prof_PriceDA.Data[8325] := 0.1475928;
   Prof_PriceDA.Data[8326] := 0.1475928;
   Prof_PriceDA.Data[8327] := 0.1475928;
   Prof_PriceDA.Data[8328] := 0.1800792;
   Prof_PriceDA.Data[8329] := 0.1800792;
   Prof_PriceDA.Data[8330] := 0.1800792;
   Prof_PriceDA.Data[8331] := 0.1800792;
   Prof_PriceDA.Data[8332] := 0.1791612;
   Prof_PriceDA.Data[8333] := 0.1791612;
   Prof_PriceDA.Data[8334] := 0.1791612;
   Prof_PriceDA.Data[8335] := 0.1791612;
   Prof_PriceDA.Data[8336] := 0.1642248;
   Prof_PriceDA.Data[8337] := 0.1642248;
   Prof_PriceDA.Data[8338] := 0.1642248;
   Prof_PriceDA.Data[8339] := 0.1642248;
   Prof_PriceDA.Data[8340] := 0.139266;
   Prof_PriceDA.Data[8341] := 0.139266;
   Prof_PriceDA.Data[8342] := 0.139266;
   Prof_PriceDA.Data[8343] := 0.139266;
   Prof_PriceDA.Data[8344] := 0.1315224;
   Prof_PriceDA.Data[8345] := 0.1315224;
   Prof_PriceDA.Data[8346] := 0.1315224;
   Prof_PriceDA.Data[8347] := 0.1315224;
   Prof_PriceDA.Data[8348] := 0.1212516;
   Prof_PriceDA.Data[8349] := 0.1212516;
   Prof_PriceDA.Data[8350] := 0.1212516;
   Prof_PriceDA.Data[8351] := 0.1212516;
   Prof_PriceDA.Data[8352] := 0.1260792;
   Prof_PriceDA.Data[8353] := 0.1260792;
   Prof_PriceDA.Data[8354] := 0.1260792;
   Prof_PriceDA.Data[8355] := 0.1260792;
   Prof_PriceDA.Data[8356] := 0.1137672;
   Prof_PriceDA.Data[8357] := 0.1137672;
   Prof_PriceDA.Data[8358] := 0.1137672;
   Prof_PriceDA.Data[8359] := 0.1137672;
   Prof_PriceDA.Data[8360] := 0.1047384;
   Prof_PriceDA.Data[8361] := 0.1047384;
   Prof_PriceDA.Data[8362] := 0.1047384;
   Prof_PriceDA.Data[8363] := 0.1047384;
   Prof_PriceDA.Data[8364] := 0.1047708;
   Prof_PriceDA.Data[8365] := 0.1047708;
   Prof_PriceDA.Data[8366] := 0.1047708;
   Prof_PriceDA.Data[8367] := 0.1047708;
   Prof_PriceDA.Data[8368] := 0.1076652;
   Prof_PriceDA.Data[8369] := 0.1076652;
   Prof_PriceDA.Data[8370] := 0.1076652;
   Prof_PriceDA.Data[8371] := 0.1076652;
   Prof_PriceDA.Data[8372] := 0.1040364;
   Prof_PriceDA.Data[8373] := 0.1040364;
   Prof_PriceDA.Data[8374] := 0.1040364;
   Prof_PriceDA.Data[8375] := 0.1040364;
   Prof_PriceDA.Data[8376] := 0.0920052;
   Prof_PriceDA.Data[8377] := 0.0920052;
   Prof_PriceDA.Data[8378] := 0.0920052;
   Prof_PriceDA.Data[8379] := 0.0920052;
   Prof_PriceDA.Data[8380] := 0.1079244;
   Prof_PriceDA.Data[8381] := 0.1079244;
   Prof_PriceDA.Data[8382] := 0.1079244;
   Prof_PriceDA.Data[8383] := 0.1079244;
   Prof_PriceDA.Data[8384] := 0.102654;
   Prof_PriceDA.Data[8385] := 0.102654;
   Prof_PriceDA.Data[8386] := 0.102654;
   Prof_PriceDA.Data[8387] := 0.102654;
   Prof_PriceDA.Data[8388] := 0.0875772;
   Prof_PriceDA.Data[8389] := 0.0875772;
   Prof_PriceDA.Data[8390] := 0.0875772;
   Prof_PriceDA.Data[8391] := 0.0875772;
   Prof_PriceDA.Data[8392] := 0.0980748;
   Prof_PriceDA.Data[8393] := 0.0980748;
   Prof_PriceDA.Data[8394] := 0.0980748;
   Prof_PriceDA.Data[8395] := 0.0980748;
   Prof_PriceDA.Data[8396] := 0.101952;
   Prof_PriceDA.Data[8397] := 0.101952;
   Prof_PriceDA.Data[8398] := 0.101952;
   Prof_PriceDA.Data[8399] := 0.101952;
   Prof_PriceDA.Data[8400] := 0.0973728;
   Prof_PriceDA.Data[8401] := 0.0973728;
   Prof_PriceDA.Data[8402] := 0.0973728;
   Prof_PriceDA.Data[8403] := 0.0973728;
   Prof_PriceDA.Data[8404] := 0.0860328;
   Prof_PriceDA.Data[8405] := 0.0860328;
   Prof_PriceDA.Data[8406] := 0.0860328;
   Prof_PriceDA.Data[8407] := 0.0860328;
   Prof_PriceDA.Data[8408] := 0.0907416;
   Prof_PriceDA.Data[8409] := 0.0907416;
   Prof_PriceDA.Data[8410] := 0.0907416;
   Prof_PriceDA.Data[8411] := 0.0907416;
   Prof_PriceDA.Data[8412] := 0.09612;
   Prof_PriceDA.Data[8413] := 0.09612;
   Prof_PriceDA.Data[8414] := 0.09612;
   Prof_PriceDA.Data[8415] := 0.09612;
   Prof_PriceDA.Data[8416] := 0.1204956;
   Prof_PriceDA.Data[8417] := 0.1204956;
   Prof_PriceDA.Data[8418] := 0.1204956;
   Prof_PriceDA.Data[8419] := 0.1204956;
   Prof_PriceDA.Data[8420] := 0.13689;
   Prof_PriceDA.Data[8421] := 0.13689;
   Prof_PriceDA.Data[8422] := 0.13689;
   Prof_PriceDA.Data[8423] := 0.13689;
   Prof_PriceDA.Data[8424] := 0.1678644;
   Prof_PriceDA.Data[8425] := 0.1678644;
   Prof_PriceDA.Data[8426] := 0.1678644;
   Prof_PriceDA.Data[8427] := 0.1678644;
   Prof_PriceDA.Data[8428] := 0.1719684;
   Prof_PriceDA.Data[8429] := 0.1719684;
   Prof_PriceDA.Data[8430] := 0.1719684;
   Prof_PriceDA.Data[8431] := 0.1719684;
   Prof_PriceDA.Data[8432] := 0.1418472;
   Prof_PriceDA.Data[8433] := 0.1418472;
   Prof_PriceDA.Data[8434] := 0.1418472;
   Prof_PriceDA.Data[8435] := 0.1418472;
   Prof_PriceDA.Data[8436] := 0.1155708;
   Prof_PriceDA.Data[8437] := 0.1155708;
   Prof_PriceDA.Data[8438] := 0.1155708;
   Prof_PriceDA.Data[8439] := 0.1155708;
   Prof_PriceDA.Data[8440] := 0.0931284;
   Prof_PriceDA.Data[8441] := 0.0931284;
   Prof_PriceDA.Data[8442] := 0.0931284;
   Prof_PriceDA.Data[8443] := 0.0931284;
   Prof_PriceDA.Data[8444] := 0.0756324;
   Prof_PriceDA.Data[8445] := 0.0756324;
   Prof_PriceDA.Data[8446] := 0.0756324;
   Prof_PriceDA.Data[8447] := 0.0756324;
   Prof_PriceDA.Data[8448] := 0.0499284;
   Prof_PriceDA.Data[8449] := 0.0499284;
   Prof_PriceDA.Data[8450] := 0.0499284;
   Prof_PriceDA.Data[8451] := 0.0499284;
   Prof_PriceDA.Data[8452] := 0.0171504;
   Prof_PriceDA.Data[8453] := 0.0171504;
   Prof_PriceDA.Data[8454] := 0.0171504;
   Prof_PriceDA.Data[8455] := 0.0171504;
   Prof_PriceDA.Data[8456] := 0.0054972;
   Prof_PriceDA.Data[8457] := 0.0054972;
   Prof_PriceDA.Data[8458] := 0.0054972;
   Prof_PriceDA.Data[8459] := 0.0054972;
   Prof_PriceDA.Data[8460] := 0.001296;
   Prof_PriceDA.Data[8461] := 0.001296;
   Prof_PriceDA.Data[8462] := 0.001296;
   Prof_PriceDA.Data[8463] := 0.001296;
   Prof_PriceDA.Data[8464] := 9.72E-05;
   Prof_PriceDA.Data[8465] := 9.72E-05;
   Prof_PriceDA.Data[8466] := 9.72E-05;
   Prof_PriceDA.Data[8467] := 9.72E-05;
   Prof_PriceDA.Data[8468] := 0.0011016;
   Prof_PriceDA.Data[8469] := 0.0011016;
   Prof_PriceDA.Data[8470] := 0.0011016;
   Prof_PriceDA.Data[8471] := 0.0011016;
   Prof_PriceDA.Data[8472] := 0.0011772;
   Prof_PriceDA.Data[8473] := 0.0011772;
   Prof_PriceDA.Data[8474] := 0.0011772;
   Prof_PriceDA.Data[8475] := 0.0011772;
   Prof_PriceDA.Data[8476] := 0.001728;
   Prof_PriceDA.Data[8477] := 0.001728;
   Prof_PriceDA.Data[8478] := 0.001728;
   Prof_PriceDA.Data[8479] := 0.001728;
   Prof_PriceDA.Data[8480] := 0.000108;
   Prof_PriceDA.Data[8481] := 0.000108;
   Prof_PriceDA.Data[8482] := 0.000108;
   Prof_PriceDA.Data[8483] := 0.000108;
   Prof_PriceDA.Data[8484] := -0.0008856;
   Prof_PriceDA.Data[8485] := -0.0008856;
   Prof_PriceDA.Data[8486] := -0.0008856;
   Prof_PriceDA.Data[8487] := -0.0008856;
   Prof_PriceDA.Data[8488] := -0.0044712;
   Prof_PriceDA.Data[8489] := -0.0044712;
   Prof_PriceDA.Data[8490] := -0.0044712;
   Prof_PriceDA.Data[8491] := -0.0044712;
   Prof_PriceDA.Data[8492] := -0.016794;
   Prof_PriceDA.Data[8493] := -0.016794;
   Prof_PriceDA.Data[8494] := -0.016794;
   Prof_PriceDA.Data[8495] := -0.016794;
   Prof_PriceDA.Data[8496] := -0.024732;
   Prof_PriceDA.Data[8497] := -0.024732;
   Prof_PriceDA.Data[8498] := -0.024732;
   Prof_PriceDA.Data[8499] := -0.024732;
   Prof_PriceDA.Data[8500] := -0.0234252;
   Prof_PriceDA.Data[8501] := -0.0234252;
   Prof_PriceDA.Data[8502] := -0.0234252;
   Prof_PriceDA.Data[8503] := -0.0234252;
   Prof_PriceDA.Data[8504] := -0.01161;
   Prof_PriceDA.Data[8505] := -0.01161;
   Prof_PriceDA.Data[8506] := -0.01161;
   Prof_PriceDA.Data[8507] := -0.01161;
   Prof_PriceDA.Data[8508] := -0.0038664;
   Prof_PriceDA.Data[8509] := -0.0038664;
   Prof_PriceDA.Data[8510] := -0.0038664;
   Prof_PriceDA.Data[8511] := -0.0038664;
   Prof_PriceDA.Data[8512] := -0.002214;
   Prof_PriceDA.Data[8513] := -0.002214;
   Prof_PriceDA.Data[8514] := -0.002214;
   Prof_PriceDA.Data[8515] := -0.002214;
   Prof_PriceDA.Data[8516] := 0.0343872;
   Prof_PriceDA.Data[8517] := 0.0343872;
   Prof_PriceDA.Data[8518] := 0.0343872;
   Prof_PriceDA.Data[8519] := 0.0343872;
   Prof_PriceDA.Data[8520] := 0.095202;
   Prof_PriceDA.Data[8521] := 0.095202;
   Prof_PriceDA.Data[8522] := 0.095202;
   Prof_PriceDA.Data[8523] := 0.095202;
   Prof_PriceDA.Data[8524] := 0.0986472;
   Prof_PriceDA.Data[8525] := 0.0986472;
   Prof_PriceDA.Data[8526] := 0.0986472;
   Prof_PriceDA.Data[8527] := 0.0986472;
   Prof_PriceDA.Data[8528] := 0.09558;
   Prof_PriceDA.Data[8529] := 0.09558;
   Prof_PriceDA.Data[8530] := 0.09558;
   Prof_PriceDA.Data[8531] := 0.09558;
   Prof_PriceDA.Data[8532] := 0.0917568;
   Prof_PriceDA.Data[8533] := 0.0917568;
   Prof_PriceDA.Data[8534] := 0.0917568;
   Prof_PriceDA.Data[8535] := 0.0917568;
   Prof_PriceDA.Data[8536] := 0.054864;
   Prof_PriceDA.Data[8537] := 0.054864;
   Prof_PriceDA.Data[8538] := 0.054864;
   Prof_PriceDA.Data[8539] := 0.054864;
   Prof_PriceDA.Data[8540] := 0.0783216;
   Prof_PriceDA.Data[8541] := 0.0783216;
   Prof_PriceDA.Data[8542] := 0.0783216;
   Prof_PriceDA.Data[8543] := 0.0783216;
   Prof_PriceDA.Data[8544] := 0.07101;
   Prof_PriceDA.Data[8545] := 0.07101;
   Prof_PriceDA.Data[8546] := 0.07101;
   Prof_PriceDA.Data[8547] := 0.07101;
   Prof_PriceDA.Data[8548] := 0.0717876;
   Prof_PriceDA.Data[8549] := 0.0717876;
   Prof_PriceDA.Data[8550] := 0.0717876;
   Prof_PriceDA.Data[8551] := 0.0717876;
   Prof_PriceDA.Data[8552] := 0.0763452;
   Prof_PriceDA.Data[8553] := 0.0763452;
   Prof_PriceDA.Data[8554] := 0.0763452;
   Prof_PriceDA.Data[8555] := 0.0763452;
   Prof_PriceDA.Data[8556] := 0.0797256;
   Prof_PriceDA.Data[8557] := 0.0797256;
   Prof_PriceDA.Data[8558] := 0.0797256;
   Prof_PriceDA.Data[8559] := 0.0797256;
   Prof_PriceDA.Data[8560] := 0.1066068;
   Prof_PriceDA.Data[8561] := 0.1066068;
   Prof_PriceDA.Data[8562] := 0.1066068;
   Prof_PriceDA.Data[8563] := 0.1066068;
   Prof_PriceDA.Data[8564] := 0.1601424;
   Prof_PriceDA.Data[8565] := 0.1601424;
   Prof_PriceDA.Data[8566] := 0.1601424;
   Prof_PriceDA.Data[8567] := 0.1601424;
   Prof_PriceDA.Data[8568] := 0.204714;
   Prof_PriceDA.Data[8569] := 0.204714;
   Prof_PriceDA.Data[8570] := 0.204714;
   Prof_PriceDA.Data[8571] := 0.204714;
   Prof_PriceDA.Data[8572] := 0.1906092;
   Prof_PriceDA.Data[8573] := 0.1906092;
   Prof_PriceDA.Data[8574] := 0.1906092;
   Prof_PriceDA.Data[8575] := 0.1906092;
   Prof_PriceDA.Data[8576] := 0.1490832;
   Prof_PriceDA.Data[8577] := 0.1490832;
   Prof_PriceDA.Data[8578] := 0.1490832;
   Prof_PriceDA.Data[8579] := 0.1490832;
   Prof_PriceDA.Data[8580] := 0.1241892;
   Prof_PriceDA.Data[8581] := 0.1241892;
   Prof_PriceDA.Data[8582] := 0.1241892;
   Prof_PriceDA.Data[8583] := 0.1241892;
   Prof_PriceDA.Data[8584] := 0.1147284;
   Prof_PriceDA.Data[8585] := 0.1147284;
   Prof_PriceDA.Data[8586] := 0.1147284;
   Prof_PriceDA.Data[8587] := 0.1147284;
   Prof_PriceDA.Data[8588] := 0.1007532;
   Prof_PriceDA.Data[8589] := 0.1007532;
   Prof_PriceDA.Data[8590] := 0.1007532;
   Prof_PriceDA.Data[8591] := 0.1007532;
   Prof_PriceDA.Data[8592] := 0.0931068;
   Prof_PriceDA.Data[8593] := 0.0931068;
   Prof_PriceDA.Data[8594] := 0.0931068;
   Prof_PriceDA.Data[8595] := 0.0931068;
   Prof_PriceDA.Data[8596] := 0.0853848;
   Prof_PriceDA.Data[8597] := 0.0853848;
   Prof_PriceDA.Data[8598] := 0.0853848;
   Prof_PriceDA.Data[8599] := 0.0853848;
   Prof_PriceDA.Data[8600] := 0.0827388;
   Prof_PriceDA.Data[8601] := 0.0827388;
   Prof_PriceDA.Data[8602] := 0.0827388;
   Prof_PriceDA.Data[8603] := 0.0827388;
   Prof_PriceDA.Data[8604] := 0.0965304;
   Prof_PriceDA.Data[8605] := 0.0965304;
   Prof_PriceDA.Data[8606] := 0.0965304;
   Prof_PriceDA.Data[8607] := 0.0965304;
   Prof_PriceDA.Data[8608] := 0.121014;
   Prof_PriceDA.Data[8609] := 0.121014;
   Prof_PriceDA.Data[8610] := 0.121014;
   Prof_PriceDA.Data[8611] := 0.121014;
   Prof_PriceDA.Data[8612] := 0.1552932;
   Prof_PriceDA.Data[8613] := 0.1552932;
   Prof_PriceDA.Data[8614] := 0.1552932;
   Prof_PriceDA.Data[8615] := 0.1552932;
   Prof_PriceDA.Data[8616] := 0.2376432;
   Prof_PriceDA.Data[8617] := 0.2376432;
   Prof_PriceDA.Data[8618] := 0.2376432;
   Prof_PriceDA.Data[8619] := 0.2376432;
   Prof_PriceDA.Data[8620] := 0.208602;
   Prof_PriceDA.Data[8621] := 0.208602;
   Prof_PriceDA.Data[8622] := 0.208602;
   Prof_PriceDA.Data[8623] := 0.208602;
   Prof_PriceDA.Data[8624] := 0.1483272;
   Prof_PriceDA.Data[8625] := 0.1483272;
   Prof_PriceDA.Data[8626] := 0.1483272;
   Prof_PriceDA.Data[8627] := 0.1483272;
   Prof_PriceDA.Data[8628] := 0.1257552;
   Prof_PriceDA.Data[8629] := 0.1257552;
   Prof_PriceDA.Data[8630] := 0.1257552;
   Prof_PriceDA.Data[8631] := 0.1257552;
   Prof_PriceDA.Data[8632] := 0.1110024;
   Prof_PriceDA.Data[8633] := 0.1110024;
   Prof_PriceDA.Data[8634] := 0.1110024;
   Prof_PriceDA.Data[8635] := 0.1110024;
   Prof_PriceDA.Data[8636] := 0.1108188;
   Prof_PriceDA.Data[8637] := 0.1108188;
   Prof_PriceDA.Data[8638] := 0.1108188;
   Prof_PriceDA.Data[8639] := 0.1108188;
   Prof_PriceDA.Data[8640] := 0.104544;
   Prof_PriceDA.Data[8641] := 0.104544;
   Prof_PriceDA.Data[8642] := 0.104544;
   Prof_PriceDA.Data[8643] := 0.104544;
   Prof_PriceDA.Data[8644] := 0.1025028;
   Prof_PriceDA.Data[8645] := 0.1025028;
   Prof_PriceDA.Data[8646] := 0.1025028;
   Prof_PriceDA.Data[8647] := 0.1025028;
   Prof_PriceDA.Data[8648] := 0.1041228;
   Prof_PriceDA.Data[8649] := 0.1041228;
   Prof_PriceDA.Data[8650] := 0.1041228;
   Prof_PriceDA.Data[8651] := 0.1041228;
   Prof_PriceDA.Data[8652] := 0.1015848;
   Prof_PriceDA.Data[8653] := 0.1015848;
   Prof_PriceDA.Data[8654] := 0.1015848;
   Prof_PriceDA.Data[8655] := 0.1015848;
   Prof_PriceDA.Data[8656] := 0.1119852;
   Prof_PriceDA.Data[8657] := 0.1119852;
   Prof_PriceDA.Data[8658] := 0.1119852;
   Prof_PriceDA.Data[8659] := 0.1119852;
   Prof_PriceDA.Data[8660] := 0.1436616;
   Prof_PriceDA.Data[8661] := 0.1436616;
   Prof_PriceDA.Data[8662] := 0.1436616;
   Prof_PriceDA.Data[8663] := 0.1436616;
   Prof_PriceDA.Data[8664] := 0.1899504;
   Prof_PriceDA.Data[8665] := 0.1899504;
   Prof_PriceDA.Data[8666] := 0.1899504;
   Prof_PriceDA.Data[8667] := 0.1899504;
   Prof_PriceDA.Data[8668] := 0.1721196;
   Prof_PriceDA.Data[8669] := 0.1721196;
   Prof_PriceDA.Data[8670] := 0.1721196;
   Prof_PriceDA.Data[8671] := 0.1721196;
   Prof_PriceDA.Data[8672] := 0.119016;
   Prof_PriceDA.Data[8673] := 0.119016;
   Prof_PriceDA.Data[8674] := 0.119016;
   Prof_PriceDA.Data[8675] := 0.119016;
   Prof_PriceDA.Data[8676] := 0.0971784;
   Prof_PriceDA.Data[8677] := 0.0971784;
   Prof_PriceDA.Data[8678] := 0.0971784;
   Prof_PriceDA.Data[8679] := 0.0971784;
   Prof_PriceDA.Data[8680] := 0.0837324;
   Prof_PriceDA.Data[8681] := 0.0837324;
   Prof_PriceDA.Data[8682] := 0.0837324;
   Prof_PriceDA.Data[8683] := 0.0837324;
   Prof_PriceDA.Data[8684] := 0.0729216;
   Prof_PriceDA.Data[8685] := 0.0729216;
   Prof_PriceDA.Data[8686] := 0.0729216;
   Prof_PriceDA.Data[8687] := 0.0729216;
   Prof_PriceDA.Data[8688] := 0.0497988;
   Prof_PriceDA.Data[8689] := 0.0497988;
   Prof_PriceDA.Data[8690] := 0.0497988;
   Prof_PriceDA.Data[8691] := 0.0497988;
   Prof_PriceDA.Data[8692] := 0.0529308;
   Prof_PriceDA.Data[8693] := 0.0529308;
   Prof_PriceDA.Data[8694] := 0.0529308;
   Prof_PriceDA.Data[8695] := 0.0529308;
   Prof_PriceDA.Data[8696] := 0.063774;
   Prof_PriceDA.Data[8697] := 0.063774;
   Prof_PriceDA.Data[8698] := 0.063774;
   Prof_PriceDA.Data[8699] := 0.063774;
   Prof_PriceDA.Data[8700] := 0.0988956;
   Prof_PriceDA.Data[8701] := 0.0988956;
   Prof_PriceDA.Data[8702] := 0.0988956;
   Prof_PriceDA.Data[8703] := 0.0988956;
   Prof_PriceDA.Data[8704] := 0.1104732;
   Prof_PriceDA.Data[8705] := 0.1104732;
   Prof_PriceDA.Data[8706] := 0.1104732;
   Prof_PriceDA.Data[8707] := 0.1104732;
   Prof_PriceDA.Data[8708] := 0.150822;
   Prof_PriceDA.Data[8709] := 0.150822;
   Prof_PriceDA.Data[8710] := 0.150822;
   Prof_PriceDA.Data[8711] := 0.150822;
   Prof_PriceDA.Data[8712] := 0.1844424;
   Prof_PriceDA.Data[8713] := 0.1844424;
   Prof_PriceDA.Data[8714] := 0.1844424;
   Prof_PriceDA.Data[8715] := 0.1844424;
   Prof_PriceDA.Data[8716] := 0.1531656;
   Prof_PriceDA.Data[8717] := 0.1531656;
   Prof_PriceDA.Data[8718] := 0.1531656;
   Prof_PriceDA.Data[8719] := 0.1531656;
   Prof_PriceDA.Data[8720] := 0.1248264;
   Prof_PriceDA.Data[8721] := 0.1248264;
   Prof_PriceDA.Data[8722] := 0.1248264;
   Prof_PriceDA.Data[8723] := 0.1248264;
   Prof_PriceDA.Data[8724] := 0.10611;
   Prof_PriceDA.Data[8725] := 0.10611;
   Prof_PriceDA.Data[8726] := 0.10611;
   Prof_PriceDA.Data[8727] := 0.10611;
   Prof_PriceDA.Data[8728] := 0.087804;
   Prof_PriceDA.Data[8729] := 0.087804;
   Prof_PriceDA.Data[8730] := 0.087804;
   Prof_PriceDA.Data[8731] := 0.087804;
   Prof_PriceDA.Data[8732] := 0.0763884;
   Prof_PriceDA.Data[8733] := 0.0763884;
   Prof_PriceDA.Data[8734] := 0.0763884;
   Prof_PriceDA.Data[8735] := 0.0763884;
   Prof_PriceDA.Data[8736] := 0.0763884;
   Prof_PriceDA.Data[8737] := 0.0763884;
   Prof_PriceDA.Data[8738] := 0.0763884;
   Prof_PriceDA.Data[8739] := 0.0763884;
   Prof_PriceDA.Data[8740] := 0.0763236;
   Prof_PriceDA.Data[8741] := 0.0763236;
   Prof_PriceDA.Data[8742] := 0.0763236;
   Prof_PriceDA.Data[8743] := 0.0763236;
   Prof_PriceDA.Data[8744] := 0.0782244;
   Prof_PriceDA.Data[8745] := 0.0782244;
   Prof_PriceDA.Data[8746] := 0.0782244;
   Prof_PriceDA.Data[8747] := 0.0782244;
   Prof_PriceDA.Data[8748] := 0.0793692;
   Prof_PriceDA.Data[8749] := 0.0793692;
   Prof_PriceDA.Data[8750] := 0.0793692;
   Prof_PriceDA.Data[8751] := 0.0793692;
   Prof_PriceDA.Data[8752] := 0.094122;
   Prof_PriceDA.Data[8753] := 0.094122;
   Prof_PriceDA.Data[8754] := 0.094122;
   Prof_PriceDA.Data[8755] := 0.094122;
   Prof_PriceDA.Data[8756] := 0.1310364;
   Prof_PriceDA.Data[8757] := 0.1310364;
   Prof_PriceDA.Data[8758] := 0.1310364;
   Prof_PriceDA.Data[8759] := 0.1310364;
   Prof_PriceDA.Data[8760] := 0.1680912;
   Prof_PriceDA.Data[8761] := 0.1680912;
   Prof_PriceDA.Data[8762] := 0.1680912;
   Prof_PriceDA.Data[8763] := 0.1680912;
   Prof_PriceDA.Data[8764] := 0.1364364;
   Prof_PriceDA.Data[8765] := 0.1364364;
   Prof_PriceDA.Data[8766] := 0.1364364;
   Prof_PriceDA.Data[8767] := 0.1364364;
   Prof_PriceDA.Data[8768] := 0.0936684;
   Prof_PriceDA.Data[8769] := 0.0936684;
   Prof_PriceDA.Data[8770] := 0.0936684;
   Prof_PriceDA.Data[8771] := 0.0936684;
   Prof_PriceDA.Data[8772] := 0.0721872;
   Prof_PriceDA.Data[8773] := 0.0721872;
   Prof_PriceDA.Data[8774] := 0.0721872;
   Prof_PriceDA.Data[8775] := 0.0721872;
   Prof_PriceDA.Data[8776] := 0.0539784;
   Prof_PriceDA.Data[8777] := 0.0539784;
   Prof_PriceDA.Data[8778] := 0.0539784;
   Prof_PriceDA.Data[8779] := 0.0539784;
   Prof_PriceDA.Data[8780] := 0.0527688;
   Prof_PriceDA.Data[8781] := 0.0527688;
   Prof_PriceDA.Data[8782] := 0.0527688;
   Prof_PriceDA.Data[8783] := 0.0527688;
   Prof_PriceDA.Data[8784] := 0.0516456;
   Prof_PriceDA.Data[8785] := 0.0516456;
   Prof_PriceDA.Data[8786] := 0.0516456;
   Prof_PriceDA.Data[8787] := 0.0516456;
   Prof_PriceDA.Data[8788] := 0.0528228;
   Prof_PriceDA.Data[8789] := 0.0528228;
   Prof_PriceDA.Data[8790] := 0.0528228;
   Prof_PriceDA.Data[8791] := 0.0528228;
   Prof_PriceDA.Data[8792] := 0.0762696;
   Prof_PriceDA.Data[8793] := 0.0762696;
   Prof_PriceDA.Data[8794] := 0.0762696;
   Prof_PriceDA.Data[8795] := 0.0762696;
   Prof_PriceDA.Data[8796] := 0.0892836;
   Prof_PriceDA.Data[8797] := 0.0892836;
   Prof_PriceDA.Data[8798] := 0.0892836;
   Prof_PriceDA.Data[8799] := 0.0892836;
   Prof_PriceDA.Data[8800] := 0.1145448;
   Prof_PriceDA.Data[8801] := 0.1145448;
   Prof_PriceDA.Data[8802] := 0.1145448;
   Prof_PriceDA.Data[8803] := 0.1145448;
   Prof_PriceDA.Data[8804] := 0.1249668;
   Prof_PriceDA.Data[8805] := 0.1249668;
   Prof_PriceDA.Data[8806] := 0.1249668;
   Prof_PriceDA.Data[8807] := 0.1249668;
   Prof_PriceDA.Data[8808] := 0.163296;
   Prof_PriceDA.Data[8809] := 0.163296;
   Prof_PriceDA.Data[8810] := 0.163296;
   Prof_PriceDA.Data[8811] := 0.163296;
   Prof_PriceDA.Data[8812] := 0.1449576;
   Prof_PriceDA.Data[8813] := 0.1449576;
   Prof_PriceDA.Data[8814] := 0.1449576;
   Prof_PriceDA.Data[8815] := 0.1449576;
   Prof_PriceDA.Data[8816] := 0.1180116;
   Prof_PriceDA.Data[8817] := 0.1180116;
   Prof_PriceDA.Data[8818] := 0.1180116;
   Prof_PriceDA.Data[8819] := 0.1180116;
   Prof_PriceDA.Data[8820] := 0.0979236;
   Prof_PriceDA.Data[8821] := 0.0979236;
   Prof_PriceDA.Data[8822] := 0.0979236;
   Prof_PriceDA.Data[8823] := 0.0979236;
   Prof_PriceDA.Data[8824] := 0.082134;
   Prof_PriceDA.Data[8825] := 0.082134;
   Prof_PriceDA.Data[8826] := 0.082134;
   Prof_PriceDA.Data[8827] := 0.082134;
   Prof_PriceDA.Data[8828] := 0.0786024;
   Prof_PriceDA.Data[8829] := 0.0786024;
   Prof_PriceDA.Data[8830] := 0.0786024;
   Prof_PriceDA.Data[8831] := 0.0786024;
   Prof_PriceDA.Data[8832] := 0.082242;
   Prof_PriceDA.Data[8833] := 0.082242;
   Prof_PriceDA.Data[8834] := 0.082242;
   Prof_PriceDA.Data[8835] := 0.082242;
   Prof_PriceDA.Data[8836] := 0.0783216;
   Prof_PriceDA.Data[8837] := 0.0783216;
   Prof_PriceDA.Data[8838] := 0.0783216;
   Prof_PriceDA.Data[8839] := 0.0783216;
   Prof_PriceDA.Data[8840] := 0.0791316;
   Prof_PriceDA.Data[8841] := 0.0791316;
   Prof_PriceDA.Data[8842] := 0.0791316;
   Prof_PriceDA.Data[8843] := 0.0791316;
   Prof_PriceDA.Data[8844] := 0.085266;
   Prof_PriceDA.Data[8845] := 0.085266;
   Prof_PriceDA.Data[8846] := 0.085266;
   Prof_PriceDA.Data[8847] := 0.085266;
   Prof_PriceDA.Data[8848] := 0.1108404;
   Prof_PriceDA.Data[8849] := 0.1108404;
   Prof_PriceDA.Data[8850] := 0.1108404;
   Prof_PriceDA.Data[8851] := 0.1108404;
   Prof_PriceDA.Data[8852] := 0.1525068;
   Prof_PriceDA.Data[8853] := 0.1525068;
   Prof_PriceDA.Data[8854] := 0.1525068;
   Prof_PriceDA.Data[8855] := 0.1525068;
   Prof_PriceDA.Data[8856] := 0.1803168;
   Prof_PriceDA.Data[8857] := 0.1803168;
   Prof_PriceDA.Data[8858] := 0.1803168;
   Prof_PriceDA.Data[8859] := 0.1803168;
   Prof_PriceDA.Data[8860] := 0.143964;
   Prof_PriceDA.Data[8861] := 0.143964;
   Prof_PriceDA.Data[8862] := 0.143964;
   Prof_PriceDA.Data[8863] := 0.143964;
   Prof_PriceDA.Data[8864] := 0.0854388;
   Prof_PriceDA.Data[8865] := 0.0854388;
   Prof_PriceDA.Data[8866] := 0.0854388;
   Prof_PriceDA.Data[8867] := 0.0854388;
   Prof_PriceDA.Data[8868] := 0.0449388;
   Prof_PriceDA.Data[8869] := 0.0449388;
   Prof_PriceDA.Data[8870] := 0.0449388;
   Prof_PriceDA.Data[8871] := 0.0449388;
   Prof_PriceDA.Data[8872] := 0.0023436;
   Prof_PriceDA.Data[8873] := 0.0023436;
   Prof_PriceDA.Data[8874] := 0.0023436;
   Prof_PriceDA.Data[8875] := 0.0023436;
   Prof_PriceDA.Data[8876] := -5.4E-05;
   Prof_PriceDA.Data[8877] := -5.4E-05;
   Prof_PriceDA.Data[8878] := -5.4E-05;
   Prof_PriceDA.Data[8879] := -5.4E-05;
   Prof_PriceDA.Data[8880] := -0.0026676;
   Prof_PriceDA.Data[8881] := -0.0026676;
   Prof_PriceDA.Data[8882] := -0.0026676;
   Prof_PriceDA.Data[8883] := -0.0026676;
   Prof_PriceDA.Data[8884] := 7.56E-05;
   Prof_PriceDA.Data[8885] := 7.56E-05;
   Prof_PriceDA.Data[8886] := 7.56E-05;
   Prof_PriceDA.Data[8887] := 7.56E-05;
   Prof_PriceDA.Data[8888] := 0.0056268;
   Prof_PriceDA.Data[8889] := 0.0056268;
   Prof_PriceDA.Data[8890] := 0.0056268;
   Prof_PriceDA.Data[8891] := 0.0056268;
   Prof_PriceDA.Data[8892] := 0.0464508;
   Prof_PriceDA.Data[8893] := 0.0464508;
   Prof_PriceDA.Data[8894] := 0.0464508;
   Prof_PriceDA.Data[8895] := 0.0464508;
   Prof_PriceDA.Data[8896] := 0.0988416;
   Prof_PriceDA.Data[8897] := 0.0988416;
   Prof_PriceDA.Data[8898] := 0.0988416;
   Prof_PriceDA.Data[8899] := 0.0988416;
   Prof_PriceDA.Data[8900] := 0.15768;
   Prof_PriceDA.Data[8901] := 0.15768;
   Prof_PriceDA.Data[8902] := 0.15768;
   Prof_PriceDA.Data[8903] := 0.15768;
   Prof_PriceDA.Data[8904] := 0.2069928;
   Prof_PriceDA.Data[8905] := 0.2069928;
   Prof_PriceDA.Data[8906] := 0.2069928;
   Prof_PriceDA.Data[8907] := 0.2069928;
   Prof_PriceDA.Data[8908] := 0.1957824;
   Prof_PriceDA.Data[8909] := 0.1957824;
   Prof_PriceDA.Data[8910] := 0.1957824;
   Prof_PriceDA.Data[8911] := 0.1957824;
   Prof_PriceDA.Data[8912] := 0.155196;
   Prof_PriceDA.Data[8913] := 0.155196;
   Prof_PriceDA.Data[8914] := 0.155196;
   Prof_PriceDA.Data[8915] := 0.155196;
   Prof_PriceDA.Data[8916] := 0.1250748;
   Prof_PriceDA.Data[8917] := 0.1250748;
   Prof_PriceDA.Data[8918] := 0.1250748;
   Prof_PriceDA.Data[8919] := 0.1250748;
   Prof_PriceDA.Data[8920] := 0.115398;
   Prof_PriceDA.Data[8921] := 0.115398;
   Prof_PriceDA.Data[8922] := 0.115398;
   Prof_PriceDA.Data[8923] := 0.115398;
   Prof_PriceDA.Data[8924] := 0.120636;
   Prof_PriceDA.Data[8925] := 0.120636;
   Prof_PriceDA.Data[8926] := 0.120636;
   Prof_PriceDA.Data[8927] := 0.120636;
   Prof_PriceDA.Data[8928] := 0.1153656;
   Prof_PriceDA.Data[8929] := 0.1153656;
   Prof_PriceDA.Data[8930] := 0.1153656;
   Prof_PriceDA.Data[8931] := 0.1153656;
   Prof_PriceDA.Data[8932] := 0.1161432;
   Prof_PriceDA.Data[8933] := 0.1161432;
   Prof_PriceDA.Data[8934] := 0.1161432;
   Prof_PriceDA.Data[8935] := 0.1161432;
   Prof_PriceDA.Data[8936] := 0.1162404;
   Prof_PriceDA.Data[8937] := 0.1162404;
   Prof_PriceDA.Data[8938] := 0.1162404;
   Prof_PriceDA.Data[8939] := 0.1162404;
   Prof_PriceDA.Data[8940] := 0.1199124;
   Prof_PriceDA.Data[8941] := 0.1199124;
   Prof_PriceDA.Data[8942] := 0.1199124;
   Prof_PriceDA.Data[8943] := 0.1199124;
   Prof_PriceDA.Data[8944] := 0.1269432;
   Prof_PriceDA.Data[8945] := 0.1269432;
   Prof_PriceDA.Data[8946] := 0.1269432;
   Prof_PriceDA.Data[8947] := 0.1269432;
   Prof_PriceDA.Data[8948] := 0.1723032;
   Prof_PriceDA.Data[8949] := 0.1723032;
   Prof_PriceDA.Data[8950] := 0.1723032;
   Prof_PriceDA.Data[8951] := 0.1723032;
   Prof_PriceDA.Data[8952] := 0.2012256;
   Prof_PriceDA.Data[8953] := 0.2012256;
   Prof_PriceDA.Data[8954] := 0.2012256;
   Prof_PriceDA.Data[8955] := 0.2012256;
   Prof_PriceDA.Data[8956] := 0.1536516;
   Prof_PriceDA.Data[8957] := 0.1536516;
   Prof_PriceDA.Data[8958] := 0.1536516;
   Prof_PriceDA.Data[8959] := 0.1536516;
   Prof_PriceDA.Data[8960] := 0.1045656;
   Prof_PriceDA.Data[8961] := 0.1045656;
   Prof_PriceDA.Data[8962] := 0.1045656;
   Prof_PriceDA.Data[8963] := 0.1045656;
   Prof_PriceDA.Data[8964] := 0.0711828;
   Prof_PriceDA.Data[8965] := 0.0711828;
   Prof_PriceDA.Data[8966] := 0.0711828;
   Prof_PriceDA.Data[8967] := 0.0711828;
   Prof_PriceDA.Data[8968] := 0.0084456;
   Prof_PriceDA.Data[8969] := 0.0084456;
   Prof_PriceDA.Data[8970] := 0.0084456;
   Prof_PriceDA.Data[8971] := 0.0084456;
   Prof_PriceDA.Data[8972] := 0.0;
   Prof_PriceDA.Data[8973] := 0.0;
   Prof_PriceDA.Data[8974] := 0.0;
   Prof_PriceDA.Data[8975] := 0.0;
   Prof_PriceDA.Data[8976] := -0.000864;
   Prof_PriceDA.Data[8977] := -0.000864;
   Prof_PriceDA.Data[8978] := -0.000864;
   Prof_PriceDA.Data[8979] := -0.000864;
   Prof_PriceDA.Data[8980] := -0.000702;
   Prof_PriceDA.Data[8981] := -0.000702;
   Prof_PriceDA.Data[8982] := -0.000702;
   Prof_PriceDA.Data[8983] := -0.000702;
   Prof_PriceDA.Data[8984] := 0.0011124;
   Prof_PriceDA.Data[8985] := 0.0011124;
   Prof_PriceDA.Data[8986] := 0.0011124;
   Prof_PriceDA.Data[8987] := 0.0011124;
   Prof_PriceDA.Data[8988] := 0.0440208;
   Prof_PriceDA.Data[8989] := 0.0440208;
   Prof_PriceDA.Data[8990] := 0.0440208;
   Prof_PriceDA.Data[8991] := 0.0440208;
   Prof_PriceDA.Data[8992] := 0.1187568;
   Prof_PriceDA.Data[8993] := 0.1187568;
   Prof_PriceDA.Data[8994] := 0.1187568;
   Prof_PriceDA.Data[8995] := 0.1187568;
   Prof_PriceDA.Data[8996] := 0.144018;
   Prof_PriceDA.Data[8997] := 0.144018;
   Prof_PriceDA.Data[8998] := 0.144018;
   Prof_PriceDA.Data[8999] := 0.144018;
   Prof_PriceDA.Data[9000] := 0.1943892;
   Prof_PriceDA.Data[9001] := 0.1943892;
   Prof_PriceDA.Data[9002] := 0.1943892;
   Prof_PriceDA.Data[9003] := 0.1943892;
   Prof_PriceDA.Data[9004] := 0.1816884;
   Prof_PriceDA.Data[9005] := 0.1816884;
   Prof_PriceDA.Data[9006] := 0.1816884;
   Prof_PriceDA.Data[9007] := 0.1816884;
   Prof_PriceDA.Data[9008] := 0.1463508;
   Prof_PriceDA.Data[9009] := 0.1463508;
   Prof_PriceDA.Data[9010] := 0.1463508;
   Prof_PriceDA.Data[9011] := 0.1463508;
   Prof_PriceDA.Data[9012] := 0.1414044;
   Prof_PriceDA.Data[9013] := 0.1414044;
   Prof_PriceDA.Data[9014] := 0.1414044;
   Prof_PriceDA.Data[9015] := 0.1414044;
   Prof_PriceDA.Data[9016] := 0.120312;
   Prof_PriceDA.Data[9017] := 0.120312;
   Prof_PriceDA.Data[9018] := 0.120312;
   Prof_PriceDA.Data[9019] := 0.120312;
   Prof_PriceDA.Data[9020] := 0.1343952;
   Prof_PriceDA.Data[9021] := 0.1343952;
   Prof_PriceDA.Data[9022] := 0.1343952;
   Prof_PriceDA.Data[9023] := 0.1343952;
   Prof_PriceDA.Data[9024] := 0.121824;
   Prof_PriceDA.Data[9025] := 0.121824;
   Prof_PriceDA.Data[9026] := 0.121824;
   Prof_PriceDA.Data[9027] := 0.121824;
   Prof_PriceDA.Data[9028] := 0.117882;
   Prof_PriceDA.Data[9029] := 0.117882;
   Prof_PriceDA.Data[9030] := 0.117882;
   Prof_PriceDA.Data[9031] := 0.117882;
   Prof_PriceDA.Data[9032] := 0.1172556;
   Prof_PriceDA.Data[9033] := 0.1172556;
   Prof_PriceDA.Data[9034] := 0.1172556;
   Prof_PriceDA.Data[9035] := 0.1172556;
   Prof_PriceDA.Data[9036] := 0.1168344;
   Prof_PriceDA.Data[9037] := 0.1168344;
   Prof_PriceDA.Data[9038] := 0.1168344;
   Prof_PriceDA.Data[9039] := 0.1168344;
   Prof_PriceDA.Data[9040] := 0.1170072;
   Prof_PriceDA.Data[9041] := 0.1170072;
   Prof_PriceDA.Data[9042] := 0.1170072;
   Prof_PriceDA.Data[9043] := 0.1170072;
   Prof_PriceDA.Data[9044] := 0.1300752;
   Prof_PriceDA.Data[9045] := 0.1300752;
   Prof_PriceDA.Data[9046] := 0.1300752;
   Prof_PriceDA.Data[9047] := 0.1300752;
   Prof_PriceDA.Data[9048] := 0.1264248;
   Prof_PriceDA.Data[9049] := 0.1264248;
   Prof_PriceDA.Data[9050] := 0.1264248;
   Prof_PriceDA.Data[9051] := 0.1264248;
   Prof_PriceDA.Data[9052] := 0.1114776;
   Prof_PriceDA.Data[9053] := 0.1114776;
   Prof_PriceDA.Data[9054] := 0.1114776;
   Prof_PriceDA.Data[9055] := 0.1114776;
   Prof_PriceDA.Data[9056] := 0.0626724;
   Prof_PriceDA.Data[9057] := 0.0626724;
   Prof_PriceDA.Data[9058] := 0.0626724;
   Prof_PriceDA.Data[9059] := 0.0626724;
   Prof_PriceDA.Data[9060] := 0.0007128;
   Prof_PriceDA.Data[9061] := 0.0007128;
   Prof_PriceDA.Data[9062] := 0.0007128;
   Prof_PriceDA.Data[9063] := 0.0007128;
   Prof_PriceDA.Data[9064] := -0.0008424;
   Prof_PriceDA.Data[9065] := -0.0008424;
   Prof_PriceDA.Data[9066] := -0.0008424;
   Prof_PriceDA.Data[9067] := -0.0008424;
   Prof_PriceDA.Data[9068] := -0.0193104;
   Prof_PriceDA.Data[9069] := -0.0193104;
   Prof_PriceDA.Data[9070] := -0.0193104;
   Prof_PriceDA.Data[9071] := -0.0193104;
   Prof_PriceDA.Data[9072] := -0.0406296;
   Prof_PriceDA.Data[9073] := -0.0406296;
   Prof_PriceDA.Data[9074] := -0.0406296;
   Prof_PriceDA.Data[9075] := -0.0406296;
   Prof_PriceDA.Data[9076] := -0.0391392;
   Prof_PriceDA.Data[9077] := -0.0391392;
   Prof_PriceDA.Data[9078] := -0.0391392;
   Prof_PriceDA.Data[9079] := -0.0391392;
   Prof_PriceDA.Data[9080] := -0.027378;
   Prof_PriceDA.Data[9081] := -0.027378;
   Prof_PriceDA.Data[9082] := -0.027378;
   Prof_PriceDA.Data[9083] := -0.027378;
   Prof_PriceDA.Data[9084] := 0.0044712;
   Prof_PriceDA.Data[9085] := 0.0044712;
   Prof_PriceDA.Data[9086] := 0.0044712;
   Prof_PriceDA.Data[9087] := 0.0044712;
   Prof_PriceDA.Data[9088] := 0.0357912;
   Prof_PriceDA.Data[9089] := 0.0357912;
   Prof_PriceDA.Data[9090] := 0.0357912;
   Prof_PriceDA.Data[9091] := 0.0357912;
   Prof_PriceDA.Data[9092] := 0.0894132;
   Prof_PriceDA.Data[9093] := 0.0894132;
   Prof_PriceDA.Data[9094] := 0.0894132;
   Prof_PriceDA.Data[9095] := 0.0894132;
   Prof_PriceDA.Data[9096] := 0.1547208;
   Prof_PriceDA.Data[9097] := 0.1547208;
   Prof_PriceDA.Data[9098] := 0.1547208;
   Prof_PriceDA.Data[9099] := 0.1547208;
   Prof_PriceDA.Data[9100] := 0.1366092;
   Prof_PriceDA.Data[9101] := 0.1366092;
   Prof_PriceDA.Data[9102] := 0.1366092;
   Prof_PriceDA.Data[9103] := 0.1366092;
   Prof_PriceDA.Data[9104] := 0.1053432;
   Prof_PriceDA.Data[9105] := 0.1053432;
   Prof_PriceDA.Data[9106] := 0.1053432;
   Prof_PriceDA.Data[9107] := 0.1053432;
   Prof_PriceDA.Data[9108] := 0.0853092;
   Prof_PriceDA.Data[9109] := 0.0853092;
   Prof_PriceDA.Data[9110] := 0.0853092;
   Prof_PriceDA.Data[9111] := 0.0853092;
   Prof_PriceDA.Data[9112] := 0.07425;
   Prof_PriceDA.Data[9113] := 0.07425;
   Prof_PriceDA.Data[9114] := 0.07425;
   Prof_PriceDA.Data[9115] := 0.07425;
   Prof_PriceDA.Data[9116] := 0.076086;
   Prof_PriceDA.Data[9117] := 0.076086;
   Prof_PriceDA.Data[9118] := 0.076086;
   Prof_PriceDA.Data[9119] := 0.076086;
   Prof_PriceDA.Data[9120] := 0.0674892;
   Prof_PriceDA.Data[9121] := 0.0674892;
   Prof_PriceDA.Data[9122] := 0.0674892;
   Prof_PriceDA.Data[9123] := 0.0674892;
   Prof_PriceDA.Data[9124] := 0.06993;
   Prof_PriceDA.Data[9125] := 0.06993;
   Prof_PriceDA.Data[9126] := 0.06993;
   Prof_PriceDA.Data[9127] := 0.06993;
   Prof_PriceDA.Data[9128] := 0.0769716;
   Prof_PriceDA.Data[9129] := 0.0769716;
   Prof_PriceDA.Data[9130] := 0.0769716;
   Prof_PriceDA.Data[9131] := 0.0769716;
   Prof_PriceDA.Data[9132] := 0.0790452;
   Prof_PriceDA.Data[9133] := 0.0790452;
   Prof_PriceDA.Data[9134] := 0.0790452;
   Prof_PriceDA.Data[9135] := 0.0790452;
   Prof_PriceDA.Data[9136] := 0.0877068;
   Prof_PriceDA.Data[9137] := 0.0877068;
   Prof_PriceDA.Data[9138] := 0.0877068;
   Prof_PriceDA.Data[9139] := 0.0877068;
   Prof_PriceDA.Data[9140] := 0.086724;
   Prof_PriceDA.Data[9141] := 0.086724;
   Prof_PriceDA.Data[9142] := 0.086724;
   Prof_PriceDA.Data[9143] := 0.086724;
   Prof_PriceDA.Data[9144] := 0.088398;
   Prof_PriceDA.Data[9145] := 0.088398;
   Prof_PriceDA.Data[9146] := 0.088398;
   Prof_PriceDA.Data[9147] := 0.088398;
   Prof_PriceDA.Data[9148] := 0.0452952;
   Prof_PriceDA.Data[9149] := 0.0452952;
   Prof_PriceDA.Data[9150] := 0.0452952;
   Prof_PriceDA.Data[9151] := 0.0452952;
   Prof_PriceDA.Data[9152] := 0.000108;
   Prof_PriceDA.Data[9153] := 0.000108;
   Prof_PriceDA.Data[9154] := 0.000108;
   Prof_PriceDA.Data[9155] := 0.000108;
   Prof_PriceDA.Data[9156] := -0.0017064;
   Prof_PriceDA.Data[9157] := -0.0017064;
   Prof_PriceDA.Data[9158] := -0.0017064;
   Prof_PriceDA.Data[9159] := -0.0017064;
   Prof_PriceDA.Data[9160] := -0.0238572;
   Prof_PriceDA.Data[9161] := -0.0238572;
   Prof_PriceDA.Data[9162] := -0.0238572;
   Prof_PriceDA.Data[9163] := -0.0238572;
   Prof_PriceDA.Data[9164] := -0.053676;
   Prof_PriceDA.Data[9165] := -0.053676;
   Prof_PriceDA.Data[9166] := -0.053676;
   Prof_PriceDA.Data[9167] := -0.053676;
   Prof_PriceDA.Data[9168] := -0.078732;
   Prof_PriceDA.Data[9169] := -0.078732;
   Prof_PriceDA.Data[9170] := -0.078732;
   Prof_PriceDA.Data[9171] := -0.078732;
   Prof_PriceDA.Data[9172] := -0.0623376;
   Prof_PriceDA.Data[9173] := -0.0623376;
   Prof_PriceDA.Data[9174] := -0.0623376;
   Prof_PriceDA.Data[9175] := -0.0623376;
   Prof_PriceDA.Data[9176] := -0.0312228;
   Prof_PriceDA.Data[9177] := -0.0312228;
   Prof_PriceDA.Data[9178] := -0.0312228;
   Prof_PriceDA.Data[9179] := -0.0312228;
   Prof_PriceDA.Data[9180] := -0.0057672;
   Prof_PriceDA.Data[9181] := -0.0057672;
   Prof_PriceDA.Data[9182] := -0.0057672;
   Prof_PriceDA.Data[9183] := -0.0057672;
   Prof_PriceDA.Data[9184] := 0.0648432;
   Prof_PriceDA.Data[9185] := 0.0648432;
   Prof_PriceDA.Data[9186] := 0.0648432;
   Prof_PriceDA.Data[9187] := 0.0648432;
   Prof_PriceDA.Data[9188] := 0.147474;
   Prof_PriceDA.Data[9189] := 0.147474;
   Prof_PriceDA.Data[9190] := 0.147474;
   Prof_PriceDA.Data[9191] := 0.147474;
   Prof_PriceDA.Data[9192] := 0.1614384;
   Prof_PriceDA.Data[9193] := 0.1614384;
   Prof_PriceDA.Data[9194] := 0.1614384;
   Prof_PriceDA.Data[9195] := 0.1614384;
   Prof_PriceDA.Data[9196] := 0.1543968;
   Prof_PriceDA.Data[9197] := 0.1543968;
   Prof_PriceDA.Data[9198] := 0.1543968;
   Prof_PriceDA.Data[9199] := 0.1543968;
   Prof_PriceDA.Data[9200] := 0.1360368;
   Prof_PriceDA.Data[9201] := 0.1360368;
   Prof_PriceDA.Data[9202] := 0.1360368;
   Prof_PriceDA.Data[9203] := 0.1360368;
   Prof_PriceDA.Data[9204] := 0.1243404;
   Prof_PriceDA.Data[9205] := 0.1243404;
   Prof_PriceDA.Data[9206] := 0.1243404;
   Prof_PriceDA.Data[9207] := 0.1243404;
   Prof_PriceDA.Data[9208] := 0.1108836;
   Prof_PriceDA.Data[9209] := 0.1108836;
   Prof_PriceDA.Data[9210] := 0.1108836;
   Prof_PriceDA.Data[9211] := 0.1108836;
   Prof_PriceDA.Data[9212] := 0.0975888;
   Prof_PriceDA.Data[9213] := 0.0975888;
   Prof_PriceDA.Data[9214] := 0.0975888;
   Prof_PriceDA.Data[9215] := 0.0975888;
   Prof_PriceDA.Data[9216] := 0.0961956;
   Prof_PriceDA.Data[9217] := 0.0961956;
   Prof_PriceDA.Data[9218] := 0.0961956;
   Prof_PriceDA.Data[9219] := 0.0961956;
   Prof_PriceDA.Data[9220] := 0.0922104;
   Prof_PriceDA.Data[9221] := 0.0922104;
   Prof_PriceDA.Data[9222] := 0.0922104;
   Prof_PriceDA.Data[9223] := 0.0922104;
   Prof_PriceDA.Data[9224] := 0.0947268;
   Prof_PriceDA.Data[9225] := 0.0947268;
   Prof_PriceDA.Data[9226] := 0.0947268;
   Prof_PriceDA.Data[9227] := 0.0947268;
   Prof_PriceDA.Data[9228] := 0.0965844;
   Prof_PriceDA.Data[9229] := 0.0965844;
   Prof_PriceDA.Data[9230] := 0.0965844;
   Prof_PriceDA.Data[9231] := 0.0965844;
   Prof_PriceDA.Data[9232] := 0.1113912;
   Prof_PriceDA.Data[9233] := 0.1113912;
   Prof_PriceDA.Data[9234] := 0.1113912;
   Prof_PriceDA.Data[9235] := 0.1113912;
   Prof_PriceDA.Data[9236] := 0.1432188;
   Prof_PriceDA.Data[9237] := 0.1432188;
   Prof_PriceDA.Data[9238] := 0.1432188;
   Prof_PriceDA.Data[9239] := 0.1432188;
   Prof_PriceDA.Data[9240] := 0.1895832;
   Prof_PriceDA.Data[9241] := 0.1895832;
   Prof_PriceDA.Data[9242] := 0.1895832;
   Prof_PriceDA.Data[9243] := 0.1895832;
   Prof_PriceDA.Data[9244] := 0.1559088;
   Prof_PriceDA.Data[9245] := 0.1559088;
   Prof_PriceDA.Data[9246] := 0.1559088;
   Prof_PriceDA.Data[9247] := 0.1559088;
   Prof_PriceDA.Data[9248] := 0.1177956;
   Prof_PriceDA.Data[9249] := 0.1177956;
   Prof_PriceDA.Data[9250] := 0.1177956;
   Prof_PriceDA.Data[9251] := 0.1177956;
   Prof_PriceDA.Data[9252] := 0.091692;
   Prof_PriceDA.Data[9253] := 0.091692;
   Prof_PriceDA.Data[9254] := 0.091692;
   Prof_PriceDA.Data[9255] := 0.091692;
   Prof_PriceDA.Data[9256] := 0.069714;
   Prof_PriceDA.Data[9257] := 0.069714;
   Prof_PriceDA.Data[9258] := 0.069714;
   Prof_PriceDA.Data[9259] := 0.069714;
   Prof_PriceDA.Data[9260] := 0.044496;
   Prof_PriceDA.Data[9261] := 0.044496;
   Prof_PriceDA.Data[9262] := 0.044496;
   Prof_PriceDA.Data[9263] := 0.044496;
   Prof_PriceDA.Data[9264] := 0.0462132;
   Prof_PriceDA.Data[9265] := 0.0462132;
   Prof_PriceDA.Data[9266] := 0.0462132;
   Prof_PriceDA.Data[9267] := 0.0462132;
   Prof_PriceDA.Data[9268] := 0.0648108;
   Prof_PriceDA.Data[9269] := 0.0648108;
   Prof_PriceDA.Data[9270] := 0.0648108;
   Prof_PriceDA.Data[9271] := 0.0648108;
   Prof_PriceDA.Data[9272] := 0.0874584;
   Prof_PriceDA.Data[9273] := 0.0874584;
   Prof_PriceDA.Data[9274] := 0.0874584;
   Prof_PriceDA.Data[9275] := 0.0874584;
   Prof_PriceDA.Data[9276] := 0.1036692;
   Prof_PriceDA.Data[9277] := 0.1036692;
   Prof_PriceDA.Data[9278] := 0.1036692;
   Prof_PriceDA.Data[9279] := 0.1036692;
   Prof_PriceDA.Data[9280] := 0.1245888;
   Prof_PriceDA.Data[9281] := 0.1245888;
   Prof_PriceDA.Data[9282] := 0.1245888;
   Prof_PriceDA.Data[9283] := 0.1245888;
   Prof_PriceDA.Data[9284] := 0.1679184;
   Prof_PriceDA.Data[9285] := 0.1679184;
   Prof_PriceDA.Data[9286] := 0.1679184;
   Prof_PriceDA.Data[9287] := 0.1679184;
   Prof_PriceDA.Data[9288] := 0.1964952;
   Prof_PriceDA.Data[9289] := 0.1964952;
   Prof_PriceDA.Data[9290] := 0.1964952;
   Prof_PriceDA.Data[9291] := 0.1964952;
   Prof_PriceDA.Data[9292] := 0.199206;
   Prof_PriceDA.Data[9293] := 0.199206;
   Prof_PriceDA.Data[9294] := 0.199206;
   Prof_PriceDA.Data[9295] := 0.199206;
   Prof_PriceDA.Data[9296] := 0.1556388;
   Prof_PriceDA.Data[9297] := 0.1556388;
   Prof_PriceDA.Data[9298] := 0.1556388;
   Prof_PriceDA.Data[9299] := 0.1556388;
   Prof_PriceDA.Data[9300] := 0.1374732;
   Prof_PriceDA.Data[9301] := 0.1374732;
   Prof_PriceDA.Data[9302] := 0.1374732;
   Prof_PriceDA.Data[9303] := 0.1374732;
   Prof_PriceDA.Data[9304] := 0.1198044;
   Prof_PriceDA.Data[9305] := 0.1198044;
   Prof_PriceDA.Data[9306] := 0.1198044;
   Prof_PriceDA.Data[9307] := 0.1198044;
   Prof_PriceDA.Data[9308] := 0.1027512;
   Prof_PriceDA.Data[9309] := 0.1027512;
   Prof_PriceDA.Data[9310] := 0.1027512;
   Prof_PriceDA.Data[9311] := 0.1027512;
   Prof_PriceDA.Data[9312] := 0.0974592;
   Prof_PriceDA.Data[9313] := 0.0974592;
   Prof_PriceDA.Data[9314] := 0.0974592;
   Prof_PriceDA.Data[9315] := 0.0974592;
   Prof_PriceDA.Data[9316] := 0.0986472;
   Prof_PriceDA.Data[9317] := 0.0986472;
   Prof_PriceDA.Data[9318] := 0.0986472;
   Prof_PriceDA.Data[9319] := 0.0986472;
   Prof_PriceDA.Data[9320] := 0.1008504;
   Prof_PriceDA.Data[9321] := 0.1008504;
   Prof_PriceDA.Data[9322] := 0.1008504;
   Prof_PriceDA.Data[9323] := 0.1008504;
   Prof_PriceDA.Data[9324] := 0.1032156;
   Prof_PriceDA.Data[9325] := 0.1032156;
   Prof_PriceDA.Data[9326] := 0.1032156;
   Prof_PriceDA.Data[9327] := 0.1032156;
   Prof_PriceDA.Data[9328] := 0.1205712;
   Prof_PriceDA.Data[9329] := 0.1205712;
   Prof_PriceDA.Data[9330] := 0.1205712;
   Prof_PriceDA.Data[9331] := 0.1205712;
   Prof_PriceDA.Data[9332] := 0.1641816;
   Prof_PriceDA.Data[9333] := 0.1641816;
   Prof_PriceDA.Data[9334] := 0.1641816;
   Prof_PriceDA.Data[9335] := 0.1641816;
   Prof_PriceDA.Data[9336] := 0.193914;
   Prof_PriceDA.Data[9337] := 0.193914;
   Prof_PriceDA.Data[9338] := 0.193914;
   Prof_PriceDA.Data[9339] := 0.193914;
   Prof_PriceDA.Data[9340] := 0.1477116;
   Prof_PriceDA.Data[9341] := 0.1477116;
   Prof_PriceDA.Data[9342] := 0.1477116;
   Prof_PriceDA.Data[9343] := 0.1477116;
   Prof_PriceDA.Data[9344] := 0.0986256;
   Prof_PriceDA.Data[9345] := 0.0986256;
   Prof_PriceDA.Data[9346] := 0.0986256;
   Prof_PriceDA.Data[9347] := 0.0986256;
   Prof_PriceDA.Data[9348] := 0.0863892;
   Prof_PriceDA.Data[9349] := 0.0863892;
   Prof_PriceDA.Data[9350] := 0.0863892;
   Prof_PriceDA.Data[9351] := 0.0863892;
   Prof_PriceDA.Data[9352] := 0.0829656;
   Prof_PriceDA.Data[9353] := 0.0829656;
   Prof_PriceDA.Data[9354] := 0.0829656;
   Prof_PriceDA.Data[9355] := 0.0829656;
   Prof_PriceDA.Data[9356] := 0.0634176;
   Prof_PriceDA.Data[9357] := 0.0634176;
   Prof_PriceDA.Data[9358] := 0.0634176;
   Prof_PriceDA.Data[9359] := 0.0634176;
   Prof_PriceDA.Data[9360] := 0.058482;
   Prof_PriceDA.Data[9361] := 0.058482;
   Prof_PriceDA.Data[9362] := 0.058482;
   Prof_PriceDA.Data[9363] := 0.058482;
   Prof_PriceDA.Data[9364] := 0.0728784;
   Prof_PriceDA.Data[9365] := 0.0728784;
   Prof_PriceDA.Data[9366] := 0.0728784;
   Prof_PriceDA.Data[9367] := 0.0728784;
   Prof_PriceDA.Data[9368] := 0.0916488;
   Prof_PriceDA.Data[9369] := 0.0916488;
   Prof_PriceDA.Data[9370] := 0.0916488;
   Prof_PriceDA.Data[9371] := 0.0916488;
   Prof_PriceDA.Data[9372] := 0.1005912;
   Prof_PriceDA.Data[9373] := 0.1005912;
   Prof_PriceDA.Data[9374] := 0.1005912;
   Prof_PriceDA.Data[9375] := 0.1005912;
   Prof_PriceDA.Data[9376] := 0.110322;
   Prof_PriceDA.Data[9377] := 0.110322;
   Prof_PriceDA.Data[9378] := 0.110322;
   Prof_PriceDA.Data[9379] := 0.110322;
   Prof_PriceDA.Data[9380] := 0.173988;
   Prof_PriceDA.Data[9381] := 0.173988;
   Prof_PriceDA.Data[9382] := 0.173988;
   Prof_PriceDA.Data[9383] := 0.173988;
   Prof_PriceDA.Data[9384] := 0.2445012;
   Prof_PriceDA.Data[9385] := 0.2445012;
   Prof_PriceDA.Data[9386] := 0.2445012;
   Prof_PriceDA.Data[9387] := 0.2445012;
   Prof_PriceDA.Data[9388] := 0.2341332;
   Prof_PriceDA.Data[9389] := 0.2341332;
   Prof_PriceDA.Data[9390] := 0.2341332;
   Prof_PriceDA.Data[9391] := 0.2341332;
   Prof_PriceDA.Data[9392] := 0.1611684;
   Prof_PriceDA.Data[9393] := 0.1611684;
   Prof_PriceDA.Data[9394] := 0.1611684;
   Prof_PriceDA.Data[9395] := 0.1611684;
   Prof_PriceDA.Data[9396] := 0.134622;
   Prof_PriceDA.Data[9397] := 0.134622;
   Prof_PriceDA.Data[9398] := 0.134622;
   Prof_PriceDA.Data[9399] := 0.134622;
   Prof_PriceDA.Data[9400] := 0.119988;
   Prof_PriceDA.Data[9401] := 0.119988;
   Prof_PriceDA.Data[9402] := 0.119988;
   Prof_PriceDA.Data[9403] := 0.119988;
   Prof_PriceDA.Data[9404] := 0.1241676;
   Prof_PriceDA.Data[9405] := 0.1241676;
   Prof_PriceDA.Data[9406] := 0.1241676;
   Prof_PriceDA.Data[9407] := 0.1241676;
   Prof_PriceDA.Data[9408] := 0.1159272;
   Prof_PriceDA.Data[9409] := 0.1159272;
   Prof_PriceDA.Data[9410] := 0.1159272;
   Prof_PriceDA.Data[9411] := 0.1159272;
   Prof_PriceDA.Data[9412] := 0.1125792;
   Prof_PriceDA.Data[9413] := 0.1125792;
   Prof_PriceDA.Data[9414] := 0.1125792;
   Prof_PriceDA.Data[9415] := 0.1125792;
   Prof_PriceDA.Data[9416] := 0.1121364;
   Prof_PriceDA.Data[9417] := 0.1121364;
   Prof_PriceDA.Data[9418] := 0.1121364;
   Prof_PriceDA.Data[9419] := 0.1121364;
   Prof_PriceDA.Data[9420] := 0.1148688;
   Prof_PriceDA.Data[9421] := 0.1148688;
   Prof_PriceDA.Data[9422] := 0.1148688;
   Prof_PriceDA.Data[9423] := 0.1148688;
   Prof_PriceDA.Data[9424] := 0.1344708;
   Prof_PriceDA.Data[9425] := 0.1344708;
   Prof_PriceDA.Data[9426] := 0.1344708;
   Prof_PriceDA.Data[9427] := 0.1344708;
   Prof_PriceDA.Data[9428] := 0.1790208;
   Prof_PriceDA.Data[9429] := 0.1790208;
   Prof_PriceDA.Data[9430] := 0.1790208;
   Prof_PriceDA.Data[9431] := 0.1790208;
   Prof_PriceDA.Data[9432] := 0.1892376;
   Prof_PriceDA.Data[9433] := 0.1892376;
   Prof_PriceDA.Data[9434] := 0.1892376;
   Prof_PriceDA.Data[9435] := 0.1892376;
   Prof_PriceDA.Data[9436] := 0.1422036;
   Prof_PriceDA.Data[9437] := 0.1422036;
   Prof_PriceDA.Data[9438] := 0.1422036;
   Prof_PriceDA.Data[9439] := 0.1422036;
   Prof_PriceDA.Data[9440] := 0.1101384;
   Prof_PriceDA.Data[9441] := 0.1101384;
   Prof_PriceDA.Data[9442] := 0.1101384;
   Prof_PriceDA.Data[9443] := 0.1101384;
   Prof_PriceDA.Data[9444] := 0.0935496;
   Prof_PriceDA.Data[9445] := 0.0935496;
   Prof_PriceDA.Data[9446] := 0.0935496;
   Prof_PriceDA.Data[9447] := 0.0935496;
   Prof_PriceDA.Data[9448] := 0.0719064;
   Prof_PriceDA.Data[9449] := 0.0719064;
   Prof_PriceDA.Data[9450] := 0.0719064;
   Prof_PriceDA.Data[9451] := 0.0719064;
   Prof_PriceDA.Data[9452] := 0.0168264;
   Prof_PriceDA.Data[9453] := 0.0168264;
   Prof_PriceDA.Data[9454] := 0.0168264;
   Prof_PriceDA.Data[9455] := 0.0168264;
   Prof_PriceDA.Data[9456] := 0.0208332;
   Prof_PriceDA.Data[9457] := 0.0208332;
   Prof_PriceDA.Data[9458] := 0.0208332;
   Prof_PriceDA.Data[9459] := 0.0208332;
   Prof_PriceDA.Data[9460] := 0.0560736;
   Prof_PriceDA.Data[9461] := 0.0560736;
   Prof_PriceDA.Data[9462] := 0.0560736;
   Prof_PriceDA.Data[9463] := 0.0560736;
   Prof_PriceDA.Data[9464] := 0.080298;
   Prof_PriceDA.Data[9465] := 0.080298;
   Prof_PriceDA.Data[9466] := 0.080298;
   Prof_PriceDA.Data[9467] := 0.080298;
   Prof_PriceDA.Data[9468] := 0.1092204;
   Prof_PriceDA.Data[9469] := 0.1092204;
   Prof_PriceDA.Data[9470] := 0.1092204;
   Prof_PriceDA.Data[9471] := 0.1092204;
   Prof_PriceDA.Data[9472] := 0.118692;
   Prof_PriceDA.Data[9473] := 0.118692;
   Prof_PriceDA.Data[9474] := 0.118692;
   Prof_PriceDA.Data[9475] := 0.118692;
   Prof_PriceDA.Data[9476] := 0.1336284;
   Prof_PriceDA.Data[9477] := 0.1336284;
   Prof_PriceDA.Data[9478] := 0.1336284;
   Prof_PriceDA.Data[9479] := 0.1336284;
   Prof_PriceDA.Data[9480] := 0.2242944;
   Prof_PriceDA.Data[9481] := 0.2242944;
   Prof_PriceDA.Data[9482] := 0.2242944;
   Prof_PriceDA.Data[9483] := 0.2242944;
   Prof_PriceDA.Data[9484] := 0.2358504;
   Prof_PriceDA.Data[9485] := 0.2358504;
   Prof_PriceDA.Data[9486] := 0.2358504;
   Prof_PriceDA.Data[9487] := 0.2358504;
   Prof_PriceDA.Data[9488] := 0.1809;
   Prof_PriceDA.Data[9489] := 0.1809;
   Prof_PriceDA.Data[9490] := 0.1809;
   Prof_PriceDA.Data[9491] := 0.1809;
   Prof_PriceDA.Data[9492] := 0.1442664;
   Prof_PriceDA.Data[9493] := 0.1442664;
   Prof_PriceDA.Data[9494] := 0.1442664;
   Prof_PriceDA.Data[9495] := 0.1442664;
   Prof_PriceDA.Data[9496] := 0.1234116;
   Prof_PriceDA.Data[9497] := 0.1234116;
   Prof_PriceDA.Data[9498] := 0.1234116;
   Prof_PriceDA.Data[9499] := 0.1234116;
   Prof_PriceDA.Data[9500] := 0.1139616;
   Prof_PriceDA.Data[9501] := 0.1139616;
   Prof_PriceDA.Data[9502] := 0.1139616;
   Prof_PriceDA.Data[9503] := 0.1139616;
   Prof_PriceDA.Data[9504] := 0.1056348;
   Prof_PriceDA.Data[9505] := 0.1056348;
   Prof_PriceDA.Data[9506] := 0.1056348;
   Prof_PriceDA.Data[9507] := 0.1056348;
   Prof_PriceDA.Data[9508] := 0.1038852;
   Prof_PriceDA.Data[9509] := 0.1038852;
   Prof_PriceDA.Data[9510] := 0.1038852;
   Prof_PriceDA.Data[9511] := 0.1038852;
   Prof_PriceDA.Data[9512] := 0.103032;
   Prof_PriceDA.Data[9513] := 0.103032;
   Prof_PriceDA.Data[9514] := 0.103032;
   Prof_PriceDA.Data[9515] := 0.103032;
   Prof_PriceDA.Data[9516] := 0.108972;
   Prof_PriceDA.Data[9517] := 0.108972;
   Prof_PriceDA.Data[9518] := 0.108972;
   Prof_PriceDA.Data[9519] := 0.108972;
   Prof_PriceDA.Data[9520] := 0.1207224;
   Prof_PriceDA.Data[9521] := 0.1207224;
   Prof_PriceDA.Data[9522] := 0.1207224;
   Prof_PriceDA.Data[9523] := 0.1207224;
   Prof_PriceDA.Data[9524] := 0.1610712;
   Prof_PriceDA.Data[9525] := 0.1610712;
   Prof_PriceDA.Data[9526] := 0.1610712;
   Prof_PriceDA.Data[9527] := 0.1610712;
   Prof_PriceDA.Data[9528] := 0.1946376;
   Prof_PriceDA.Data[9529] := 0.1946376;
   Prof_PriceDA.Data[9530] := 0.1946376;
   Prof_PriceDA.Data[9531] := 0.1946376;
   Prof_PriceDA.Data[9532] := 0.1502064;
   Prof_PriceDA.Data[9533] := 0.1502064;
   Prof_PriceDA.Data[9534] := 0.1502064;
   Prof_PriceDA.Data[9535] := 0.1502064;
   Prof_PriceDA.Data[9536] := 0.113184;
   Prof_PriceDA.Data[9537] := 0.113184;
   Prof_PriceDA.Data[9538] := 0.113184;
   Prof_PriceDA.Data[9539] := 0.113184;
   Prof_PriceDA.Data[9540] := 0.0890028;
   Prof_PriceDA.Data[9541] := 0.0890028;
   Prof_PriceDA.Data[9542] := 0.0890028;
   Prof_PriceDA.Data[9543] := 0.0890028;
   Prof_PriceDA.Data[9544] := 0.0739584;
   Prof_PriceDA.Data[9545] := 0.0739584;
   Prof_PriceDA.Data[9546] := 0.0739584;
   Prof_PriceDA.Data[9547] := 0.0739584;
   Prof_PriceDA.Data[9548] := 0.0424116;
   Prof_PriceDA.Data[9549] := 0.0424116;
   Prof_PriceDA.Data[9550] := 0.0424116;
   Prof_PriceDA.Data[9551] := 0.0424116;
   Prof_PriceDA.Data[9552] := 0.0027648;
   Prof_PriceDA.Data[9553] := 0.0027648;
   Prof_PriceDA.Data[9554] := 0.0027648;
   Prof_PriceDA.Data[9555] := 0.0027648;
   Prof_PriceDA.Data[9556] := 9.72E-05;
   Prof_PriceDA.Data[9557] := 9.72E-05;
   Prof_PriceDA.Data[9558] := 9.72E-05;
   Prof_PriceDA.Data[9559] := 9.72E-05;
   Prof_PriceDA.Data[9560] := 0.0023652;
   Prof_PriceDA.Data[9561] := 0.0023652;
   Prof_PriceDA.Data[9562] := 0.0023652;
   Prof_PriceDA.Data[9563] := 0.0023652;
   Prof_PriceDA.Data[9564] := 0.0735912;
   Prof_PriceDA.Data[9565] := 0.0735912;
   Prof_PriceDA.Data[9566] := 0.0735912;
   Prof_PriceDA.Data[9567] := 0.0735912;
   Prof_PriceDA.Data[9568] := 0.0892836;
   Prof_PriceDA.Data[9569] := 0.0892836;
   Prof_PriceDA.Data[9570] := 0.0892836;
   Prof_PriceDA.Data[9571] := 0.0892836;
   Prof_PriceDA.Data[9572] := 0.1238868;
   Prof_PriceDA.Data[9573] := 0.1238868;
   Prof_PriceDA.Data[9574] := 0.1238868;
   Prof_PriceDA.Data[9575] := 0.1238868;
   Prof_PriceDA.Data[9576] := 0.1767744;
   Prof_PriceDA.Data[9577] := 0.1767744;
   Prof_PriceDA.Data[9578] := 0.1767744;
   Prof_PriceDA.Data[9579] := 0.1767744;
   Prof_PriceDA.Data[9580] := 0.18414;
   Prof_PriceDA.Data[9581] := 0.18414;
   Prof_PriceDA.Data[9582] := 0.18414;
   Prof_PriceDA.Data[9583] := 0.18414;
   Prof_PriceDA.Data[9584] := 0.1397844;
   Prof_PriceDA.Data[9585] := 0.1397844;
   Prof_PriceDA.Data[9586] := 0.1397844;
   Prof_PriceDA.Data[9587] := 0.1397844;
   Prof_PriceDA.Data[9588] := 0.1205496;
   Prof_PriceDA.Data[9589] := 0.1205496;
   Prof_PriceDA.Data[9590] := 0.1205496;
   Prof_PriceDA.Data[9591] := 0.1205496;
   Prof_PriceDA.Data[9592] := 0.093258;
   Prof_PriceDA.Data[9593] := 0.093258;
   Prof_PriceDA.Data[9594] := 0.093258;
   Prof_PriceDA.Data[9595] := 0.093258;
   Prof_PriceDA.Data[9596] := 0.0891756;
   Prof_PriceDA.Data[9597] := 0.0891756;
   Prof_PriceDA.Data[9598] := 0.0891756;
   Prof_PriceDA.Data[9599] := 0.0891756;
   Prof_PriceDA.Data[9600] := 0.085266;
   Prof_PriceDA.Data[9601] := 0.085266;
   Prof_PriceDA.Data[9602] := 0.085266;
   Prof_PriceDA.Data[9603] := 0.085266;
   Prof_PriceDA.Data[9604] := 0.0749844;
   Prof_PriceDA.Data[9605] := 0.0749844;
   Prof_PriceDA.Data[9606] := 0.0749844;
   Prof_PriceDA.Data[9607] := 0.0749844;
   Prof_PriceDA.Data[9608] := 0.0763452;
   Prof_PriceDA.Data[9609] := 0.0763452;
   Prof_PriceDA.Data[9610] := 0.0763452;
   Prof_PriceDA.Data[9611] := 0.0763452;
   Prof_PriceDA.Data[9612] := 0.0837648;
   Prof_PriceDA.Data[9613] := 0.0837648;
   Prof_PriceDA.Data[9614] := 0.0837648;
   Prof_PriceDA.Data[9615] := 0.0837648;
   Prof_PriceDA.Data[9616] := 0.0936144;
   Prof_PriceDA.Data[9617] := 0.0936144;
   Prof_PriceDA.Data[9618] := 0.0936144;
   Prof_PriceDA.Data[9619] := 0.0936144;
   Prof_PriceDA.Data[9620] := 0.1195776;
   Prof_PriceDA.Data[9621] := 0.1195776;
   Prof_PriceDA.Data[9622] := 0.1195776;
   Prof_PriceDA.Data[9623] := 0.1195776;
   Prof_PriceDA.Data[9624] := 0.1210788;
   Prof_PriceDA.Data[9625] := 0.1210788;
   Prof_PriceDA.Data[9626] := 0.1210788;
   Prof_PriceDA.Data[9627] := 0.1210788;
   Prof_PriceDA.Data[9628] := 0.0954072;
   Prof_PriceDA.Data[9629] := 0.0954072;
   Prof_PriceDA.Data[9630] := 0.0954072;
   Prof_PriceDA.Data[9631] := 0.0954072;
   Prof_PriceDA.Data[9632] := 0.0687636;
   Prof_PriceDA.Data[9633] := 0.0687636;
   Prof_PriceDA.Data[9634] := 0.0687636;
   Prof_PriceDA.Data[9635] := 0.0687636;
   Prof_PriceDA.Data[9636] := 0.0160056;
   Prof_PriceDA.Data[9637] := 0.0160056;
   Prof_PriceDA.Data[9638] := 0.0160056;
   Prof_PriceDA.Data[9639] := 0.0160056;
   Prof_PriceDA.Data[9640] := 0.0003456;
   Prof_PriceDA.Data[9641] := 0.0003456;
   Prof_PriceDA.Data[9642] := 0.0003456;
   Prof_PriceDA.Data[9643] := 0.0003456;
   Prof_PriceDA.Data[9644] := -0.0001944;
   Prof_PriceDA.Data[9645] := -0.0001944;
   Prof_PriceDA.Data[9646] := -0.0001944;
   Prof_PriceDA.Data[9647] := -0.0001944;
   Prof_PriceDA.Data[9648] := -0.0003996;
   Prof_PriceDA.Data[9649] := -0.0003996;
   Prof_PriceDA.Data[9650] := -0.0003996;
   Prof_PriceDA.Data[9651] := -0.0003996;
   Prof_PriceDA.Data[9652] := -0.0012204;
   Prof_PriceDA.Data[9653] := -0.0012204;
   Prof_PriceDA.Data[9654] := -0.0012204;
   Prof_PriceDA.Data[9655] := -0.0012204;
   Prof_PriceDA.Data[9656] := -1.08E-05;
   Prof_PriceDA.Data[9657] := -1.08E-05;
   Prof_PriceDA.Data[9658] := -1.08E-05;
   Prof_PriceDA.Data[9659] := -1.08E-05;
   Prof_PriceDA.Data[9660] := 0.0644436;
   Prof_PriceDA.Data[9661] := 0.0644436;
   Prof_PriceDA.Data[9662] := 0.0644436;
   Prof_PriceDA.Data[9663] := 0.0644436;
   Prof_PriceDA.Data[9664] := 0.1005372;
   Prof_PriceDA.Data[9665] := 0.1005372;
   Prof_PriceDA.Data[9666] := 0.1005372;
   Prof_PriceDA.Data[9667] := 0.1005372;
   Prof_PriceDA.Data[9668] := 0.1495152;
   Prof_PriceDA.Data[9669] := 0.1495152;
   Prof_PriceDA.Data[9670] := 0.1495152;
   Prof_PriceDA.Data[9671] := 0.1495152;
   Prof_PriceDA.Data[9672] := 0.2005128;
   Prof_PriceDA.Data[9673] := 0.2005128;
   Prof_PriceDA.Data[9674] := 0.2005128;
   Prof_PriceDA.Data[9675] := 0.2005128;
   Prof_PriceDA.Data[9676] := 0.2052108;
   Prof_PriceDA.Data[9677] := 0.2052108;
   Prof_PriceDA.Data[9678] := 0.2052108;
   Prof_PriceDA.Data[9679] := 0.2052108;
   Prof_PriceDA.Data[9680] := 0.1707912;
   Prof_PriceDA.Data[9681] := 0.1707912;
   Prof_PriceDA.Data[9682] := 0.1707912;
   Prof_PriceDA.Data[9683] := 0.1707912;
   Prof_PriceDA.Data[9684] := 0.1496556;
   Prof_PriceDA.Data[9685] := 0.1496556;
   Prof_PriceDA.Data[9686] := 0.1496556;
   Prof_PriceDA.Data[9687] := 0.1496556;
   Prof_PriceDA.Data[9688] := 0.1200096;
   Prof_PriceDA.Data[9689] := 0.1200096;
   Prof_PriceDA.Data[9690] := 0.1200096;
   Prof_PriceDA.Data[9691] := 0.1200096;
   Prof_PriceDA.Data[9692] := 0.1212516;
   Prof_PriceDA.Data[9693] := 0.1212516;
   Prof_PriceDA.Data[9694] := 0.1212516;
   Prof_PriceDA.Data[9695] := 0.1212516;
   Prof_PriceDA.Data[9696] := 0.1176876;
   Prof_PriceDA.Data[9697] := 0.1176876;
   Prof_PriceDA.Data[9698] := 0.1176876;
   Prof_PriceDA.Data[9699] := 0.1176876;
   Prof_PriceDA.Data[9700] := 0.1135836;
   Prof_PriceDA.Data[9701] := 0.1135836;
   Prof_PriceDA.Data[9702] := 0.1135836;
   Prof_PriceDA.Data[9703] := 0.1135836;
   Prof_PriceDA.Data[9704] := 0.111672;
   Prof_PriceDA.Data[9705] := 0.111672;
   Prof_PriceDA.Data[9706] := 0.111672;
   Prof_PriceDA.Data[9707] := 0.111672;
   Prof_PriceDA.Data[9708] := 0.1126116;
   Prof_PriceDA.Data[9709] := 0.1126116;
   Prof_PriceDA.Data[9710] := 0.1126116;
   Prof_PriceDA.Data[9711] := 0.1126116;
   Prof_PriceDA.Data[9712] := 0.1131084;
   Prof_PriceDA.Data[9713] := 0.1131084;
   Prof_PriceDA.Data[9714] := 0.1131084;
   Prof_PriceDA.Data[9715] := 0.1131084;
   Prof_PriceDA.Data[9716] := 0.1209168;
   Prof_PriceDA.Data[9717] := 0.1209168;
   Prof_PriceDA.Data[9718] := 0.1209168;
   Prof_PriceDA.Data[9719] := 0.1209168;
   Prof_PriceDA.Data[9720] := 0.1166508;
   Prof_PriceDA.Data[9721] := 0.1166508;
   Prof_PriceDA.Data[9722] := 0.1166508;
   Prof_PriceDA.Data[9723] := 0.1166508;
   Prof_PriceDA.Data[9724] := 0.107244;
   Prof_PriceDA.Data[9725] := 0.107244;
   Prof_PriceDA.Data[9726] := 0.107244;
   Prof_PriceDA.Data[9727] := 0.107244;
   Prof_PriceDA.Data[9728] := 0.0751788;
   Prof_PriceDA.Data[9729] := 0.0751788;
   Prof_PriceDA.Data[9730] := 0.0751788;
   Prof_PriceDA.Data[9731] := 0.0751788;
   Prof_PriceDA.Data[9732] := 0.0218052;
   Prof_PriceDA.Data[9733] := 0.0218052;
   Prof_PriceDA.Data[9734] := 0.0218052;
   Prof_PriceDA.Data[9735] := 0.0218052;
   Prof_PriceDA.Data[9736] := 0.0;
   Prof_PriceDA.Data[9737] := 0.0;
   Prof_PriceDA.Data[9738] := 0.0;
   Prof_PriceDA.Data[9739] := 0.0;
   Prof_PriceDA.Data[9740] := -0.0082512;
   Prof_PriceDA.Data[9741] := -0.0082512;
   Prof_PriceDA.Data[9742] := -0.0082512;
   Prof_PriceDA.Data[9743] := -0.0082512;
   Prof_PriceDA.Data[9744] := -0.0096336;
   Prof_PriceDA.Data[9745] := -0.0096336;
   Prof_PriceDA.Data[9746] := -0.0096336;
   Prof_PriceDA.Data[9747] := -0.0096336;
   Prof_PriceDA.Data[9748] := -0.0296352;
   Prof_PriceDA.Data[9749] := -0.0296352;
   Prof_PriceDA.Data[9750] := -0.0296352;
   Prof_PriceDA.Data[9751] := -0.0296352;
   Prof_PriceDA.Data[9752] := -0.0058104;
   Prof_PriceDA.Data[9753] := -0.0058104;
   Prof_PriceDA.Data[9754] := -0.0058104;
   Prof_PriceDA.Data[9755] := -0.0058104;
   Prof_PriceDA.Data[9756] := 0.0024084;
   Prof_PriceDA.Data[9757] := 0.0024084;
   Prof_PriceDA.Data[9758] := 0.0024084;
   Prof_PriceDA.Data[9759] := 0.0024084;
   Prof_PriceDA.Data[9760] := 0.0930852;
   Prof_PriceDA.Data[9761] := 0.0930852;
   Prof_PriceDA.Data[9762] := 0.0930852;
   Prof_PriceDA.Data[9763] := 0.0930852;
   Prof_PriceDA.Data[9764] := 0.1310688;
   Prof_PriceDA.Data[9765] := 0.1310688;
   Prof_PriceDA.Data[9766] := 0.1310688;
   Prof_PriceDA.Data[9767] := 0.1310688;
   Prof_PriceDA.Data[9768] := 0.1958904;
   Prof_PriceDA.Data[9769] := 0.1958904;
   Prof_PriceDA.Data[9770] := 0.1958904;
   Prof_PriceDA.Data[9771] := 0.1958904;
   Prof_PriceDA.Data[9772] := 0.1957068;
   Prof_PriceDA.Data[9773] := 0.1957068;
   Prof_PriceDA.Data[9774] := 0.1957068;
   Prof_PriceDA.Data[9775] := 0.1957068;
   Prof_PriceDA.Data[9776] := 0.1428516;
   Prof_PriceDA.Data[9777] := 0.1428516;
   Prof_PriceDA.Data[9778] := 0.1428516;
   Prof_PriceDA.Data[9779] := 0.1428516;
   Prof_PriceDA.Data[9780] := 0.1317492;
   Prof_PriceDA.Data[9781] := 0.1317492;
   Prof_PriceDA.Data[9782] := 0.1317492;
   Prof_PriceDA.Data[9783] := 0.1317492;
   Prof_PriceDA.Data[9784] := 0.1090692;
   Prof_PriceDA.Data[9785] := 0.1090692;
   Prof_PriceDA.Data[9786] := 0.1090692;
   Prof_PriceDA.Data[9787] := 0.1090692;
   Prof_PriceDA.Data[9788] := 0.1047492;
   Prof_PriceDA.Data[9789] := 0.1047492;
   Prof_PriceDA.Data[9790] := 0.1047492;
   Prof_PriceDA.Data[9791] := 0.1047492;
   Prof_PriceDA.Data[9792] := 0.0844236;
   Prof_PriceDA.Data[9793] := 0.0844236;
   Prof_PriceDA.Data[9794] := 0.0844236;
   Prof_PriceDA.Data[9795] := 0.0844236;
   Prof_PriceDA.Data[9796] := 0.06723;
   Prof_PriceDA.Data[9797] := 0.06723;
   Prof_PriceDA.Data[9798] := 0.06723;
   Prof_PriceDA.Data[9799] := 0.06723;
   Prof_PriceDA.Data[9800] := 0.0808596;
   Prof_PriceDA.Data[9801] := 0.0808596;
   Prof_PriceDA.Data[9802] := 0.0808596;
   Prof_PriceDA.Data[9803] := 0.0808596;
   Prof_PriceDA.Data[9804] := 0.068904;
   Prof_PriceDA.Data[9805] := 0.068904;
   Prof_PriceDA.Data[9806] := 0.068904;
   Prof_PriceDA.Data[9807] := 0.068904;
   Prof_PriceDA.Data[9808] := 0.07047;
   Prof_PriceDA.Data[9809] := 0.07047;
   Prof_PriceDA.Data[9810] := 0.07047;
   Prof_PriceDA.Data[9811] := 0.07047;
   Prof_PriceDA.Data[9812] := 0.0669492;
   Prof_PriceDA.Data[9813] := 0.0669492;
   Prof_PriceDA.Data[9814] := 0.0669492;
   Prof_PriceDA.Data[9815] := 0.0669492;
   Prof_PriceDA.Data[9816] := 0.02997;
   Prof_PriceDA.Data[9817] := 0.02997;
   Prof_PriceDA.Data[9818] := 0.02997;
   Prof_PriceDA.Data[9819] := 0.02997;
   Prof_PriceDA.Data[9820] := 0.0145044;
   Prof_PriceDA.Data[9821] := 0.0145044;
   Prof_PriceDA.Data[9822] := 0.0145044;
   Prof_PriceDA.Data[9823] := 0.0145044;
   Prof_PriceDA.Data[9824] := 0.0091044;
   Prof_PriceDA.Data[9825] := 0.0091044;
   Prof_PriceDA.Data[9826] := 0.0091044;
   Prof_PriceDA.Data[9827] := 0.0091044;
   Prof_PriceDA.Data[9828] := 0.0;
   Prof_PriceDA.Data[9829] := 0.0;
   Prof_PriceDA.Data[9830] := 0.0;
   Prof_PriceDA.Data[9831] := 0.0;
   Prof_PriceDA.Data[9832] := -2.16E-05;
   Prof_PriceDA.Data[9833] := -2.16E-05;
   Prof_PriceDA.Data[9834] := -2.16E-05;
   Prof_PriceDA.Data[9835] := -2.16E-05;
   Prof_PriceDA.Data[9836] := -0.0039528;
   Prof_PriceDA.Data[9837] := -0.0039528;
   Prof_PriceDA.Data[9838] := -0.0039528;
   Prof_PriceDA.Data[9839] := -0.0039528;
   Prof_PriceDA.Data[9840] := -0.0203472;
   Prof_PriceDA.Data[9841] := -0.0203472;
   Prof_PriceDA.Data[9842] := -0.0203472;
   Prof_PriceDA.Data[9843] := -0.0203472;
   Prof_PriceDA.Data[9844] := -0.0274104;
   Prof_PriceDA.Data[9845] := -0.0274104;
   Prof_PriceDA.Data[9846] := -0.0274104;
   Prof_PriceDA.Data[9